(* IEC 61131-3 sources: plc-hackathon-2026/work/dump/MyController/Plc Logic/Application/Init (part 2) *)

(* ---- Init_Prof_FEC.st ---- *)
FUNCTION_BLOCK Init_Prof_FEC
VAR_INPUT
END_VAR
VAR_OUTPUT
END_VAR
VAR
END_VAR

// ---IMPL---
// Inicijalizacija GVL "Prof_FEC"
   Prof_FEC.Data[0] := 40.266;
   Prof_FEC.Data[1] := 42.108;
   Prof_FEC.Data[2] := 42.44;
   Prof_FEC.Data[3] := 43.126;
   Prof_FEC.Data[4] := 43.213;
   Prof_FEC.Data[5] := 42.172;
   Prof_FEC.Data[6] := 44.978;
   Prof_FEC.Data[7] := 44.952;
   Prof_FEC.Data[8] := 43.73;
   Prof_FEC.Data[9] := 41.671;
   Prof_FEC.Data[10] := 39.025;
   Prof_FEC.Data[11] := 43.815;
   Prof_FEC.Data[12] := 42.205;
   Prof_FEC.Data[13] := 42.881;
   Prof_FEC.Data[14] := 40.68;
   Prof_FEC.Data[15] := 39.411;
   Prof_FEC.Data[16] := 40.682;
   Prof_FEC.Data[17] := 40.404;
   Prof_FEC.Data[18] := 41.293;
   Prof_FEC.Data[19] := 41.787;
   Prof_FEC.Data[20] := 254.21;
   Prof_FEC.Data[21] := 268.75;
   Prof_FEC.Data[22] := 265.48;
   Prof_FEC.Data[23] := 296.02;
   Prof_FEC.Data[24] := 335.71;
   Prof_FEC.Data[25] := 339.43;
   Prof_FEC.Data[26] := 388.16;
   Prof_FEC.Data[27] := 433.83;
   Prof_FEC.Data[28] := 441.67;
   Prof_FEC.Data[29] := 486.31;
   Prof_FEC.Data[30] := 552.6;
   Prof_FEC.Data[31] := 544.94;
   Prof_FEC.Data[32] := 568.79;
   Prof_FEC.Data[33] := 634.46;
   Prof_FEC.Data[34] := 604.12;
   Prof_FEC.Data[35] := 630.85;
   Prof_FEC.Data[36] := 656.31;
   Prof_FEC.Data[37] := 671.59;
   Prof_FEC.Data[38] := 634.52;
   Prof_FEC.Data[39] := 653.7;
   Prof_FEC.Data[40] := 625.93;
   Prof_FEC.Data[41] := 654.27;
   Prof_FEC.Data[42] := 603.66;
   Prof_FEC.Data[43] := 590.51;
   Prof_FEC.Data[44] := 620.11;
   Prof_FEC.Data[45] := 604.33;
   Prof_FEC.Data[46] := 589.58;
   Prof_FEC.Data[47] := 638.77;
   Prof_FEC.Data[48] := 571.87;
   Prof_FEC.Data[49] := 540.78;
   Prof_FEC.Data[50] := 589.62;
   Prof_FEC.Data[51] := 576.36;
   Prof_FEC.Data[52] := 646.42;
   Prof_FEC.Data[53] := 628.77;
   Prof_FEC.Data[54] := 633.92;
   Prof_FEC.Data[55] := 671.67;
   Prof_FEC.Data[56] := 731.0;
   Prof_FEC.Data[57] := 742.29;
   Prof_FEC.Data[58] := 722.04;
   Prof_FEC.Data[59] := 711.5;
   Prof_FEC.Data[60] := 722.32;
   Prof_FEC.Data[61] := 679.4;
   Prof_FEC.Data[62] := 676.24;
   Prof_FEC.Data[63] := 745.59;
   Prof_FEC.Data[64] := 789.69;
   Prof_FEC.Data[65] := 795.4;
   Prof_FEC.Data[66] := 766.74;
   Prof_FEC.Data[67] := 673.77;
   Prof_FEC.Data[68] := 501.09;
   Prof_FEC.Data[69] := 365.1;
   Prof_FEC.Data[70] := 325.78;
   Prof_FEC.Data[71] := 293.7;
   Prof_FEC.Data[72] := 276.68;
   Prof_FEC.Data[73] := 266.17;
   Prof_FEC.Data[74] := 227.53;
   Prof_FEC.Data[75] := 256.11;
   Prof_FEC.Data[76] := 43.481;
   Prof_FEC.Data[77] := 44.002;
   Prof_FEC.Data[78] := 44.238;
   Prof_FEC.Data[79] := 43.218;
   Prof_FEC.Data[80] := 40.422;
   Prof_FEC.Data[81] := 41.151;
   Prof_FEC.Data[82] := 40.95;
   Prof_FEC.Data[83] := 41.165;
   Prof_FEC.Data[84] := 40.77;
   Prof_FEC.Data[85] := 43.799;
   Prof_FEC.Data[86] := 42.671;
   Prof_FEC.Data[87] := 43.676;
   Prof_FEC.Data[88] := 41.656;
   Prof_FEC.Data[89] := 40.912;
   Prof_FEC.Data[90] := 41.266;
   Prof_FEC.Data[91] := 39.497;
   Prof_FEC.Data[92] := 44.511;
   Prof_FEC.Data[93] := 44.6;
   Prof_FEC.Data[94] := 47.837;
   Prof_FEC.Data[95] := 45.96;
   Prof_FEC.Data[96] := 45.749;
   Prof_FEC.Data[97] := 44.326;
   Prof_FEC.Data[98] := 44.02;
   Prof_FEC.Data[99] := 43.86;
   Prof_FEC.Data[100] := 44.651;
   Prof_FEC.Data[101] := 48.206;
   Prof_FEC.Data[102] := 43.013;
   Prof_FEC.Data[103] := 45.661;
   Prof_FEC.Data[104] := 40.107;
   Prof_FEC.Data[105] := 41.976;
   Prof_FEC.Data[106] := 37.462;
   Prof_FEC.Data[107] := 40.495;
   Prof_FEC.Data[108] := 45.365;
   Prof_FEC.Data[109] := 47.462;
   Prof_FEC.Data[110] := 48.015;
   Prof_FEC.Data[111] := 48.333;
   Prof_FEC.Data[112] := 47.113;
   Prof_FEC.Data[113] := 48.016;
   Prof_FEC.Data[114] := 44.19;
   Prof_FEC.Data[115] := 45.094;
   Prof_FEC.Data[116] := 290.32;
   Prof_FEC.Data[117] := 297.39;
   Prof_FEC.Data[118] := 284.58;
   Prof_FEC.Data[119] := 325.31;
   Prof_FEC.Data[120] := 357.24;
   Prof_FEC.Data[121] := 394.59;
   Prof_FEC.Data[122] := 407.32;
   Prof_FEC.Data[123] := 458.08;
   Prof_FEC.Data[124] := 551.82;
   Prof_FEC.Data[125] := 580.15;
   Prof_FEC.Data[126] := 608.06;
   Prof_FEC.Data[127] := 578.6;
   Prof_FEC.Data[128] := 612.98;
   Prof_FEC.Data[129] := 614.51;
   Prof_FEC.Data[130] := 640.99;
   Prof_FEC.Data[131] := 677.4;
   Prof_FEC.Data[132] := 743.46;
   Prof_FEC.Data[133] := 772.07;
   Prof_FEC.Data[134] := 790.32;
   Prof_FEC.Data[135] := 764.21;
   Prof_FEC.Data[136] := 693.38;
   Prof_FEC.Data[137] := 715.42;
   Prof_FEC.Data[138] := 590.75;
   Prof_FEC.Data[139] := 678.98;
   Prof_FEC.Data[140] := 643.33;
   Prof_FEC.Data[141] := 614.71;
   Prof_FEC.Data[142] := 677.61;
   Prof_FEC.Data[143] := 646.57;
   Prof_FEC.Data[144] := 662.01;
   Prof_FEC.Data[145] := 656.44;
   Prof_FEC.Data[146] := 583.37;
   Prof_FEC.Data[147] := 664.52;
   Prof_FEC.Data[148] := 554.65;
   Prof_FEC.Data[149] := 629.64;
   Prof_FEC.Data[150] := 670.62;
   Prof_FEC.Data[151] := 596.51;
   Prof_FEC.Data[152] := 661.81;
   Prof_FEC.Data[153] := 592.39;
   Prof_FEC.Data[154] := 608.2;
   Prof_FEC.Data[155] := 668.41;
   Prof_FEC.Data[156] := 618.77;
   Prof_FEC.Data[157] := 575.67;
   Prof_FEC.Data[158] := 513.16;
   Prof_FEC.Data[159] := 598.3;
   Prof_FEC.Data[160] := 660.23;
   Prof_FEC.Data[161] := 656.71;
   Prof_FEC.Data[162] := 634.91;
   Prof_FEC.Data[163] := 512.09;
   Prof_FEC.Data[164] := 414.01;
   Prof_FEC.Data[165] := 373.69;
   Prof_FEC.Data[166] := 339.29;
   Prof_FEC.Data[167] := 286.59;
   Prof_FEC.Data[168] := 285.53;
   Prof_FEC.Data[169] := 218.56;
   Prof_FEC.Data[170] := 242.09;
   Prof_FEC.Data[171] := 257.24;
   Prof_FEC.Data[172] := 44.634;
   Prof_FEC.Data[173] := 44.75;
   Prof_FEC.Data[174] := 41.675;
   Prof_FEC.Data[175] := 49.065;
   Prof_FEC.Data[176] := 47.236;
   Prof_FEC.Data[177] := 43.529;
   Prof_FEC.Data[178] := 44.439;
   Prof_FEC.Data[179] := 44.502;
   Prof_FEC.Data[180] := 48.851;
   Prof_FEC.Data[181] := 50.0;
   Prof_FEC.Data[182] := 47.07;
   Prof_FEC.Data[183] := 44.555;
   Prof_FEC.Data[184] := 44.815;
   Prof_FEC.Data[185] := 44.276;
   Prof_FEC.Data[186] := 44.342;
   Prof_FEC.Data[187] := 43.996;
   Prof_FEC.Data[188] := 44.701;
   Prof_FEC.Data[189] := 45.391;
   Prof_FEC.Data[190] := 41.212;
   Prof_FEC.Data[191] := 44.161;
   Prof_FEC.Data[192] := 43.203;
   Prof_FEC.Data[193] := 41.683;
   Prof_FEC.Data[194] := 43.808;
   Prof_FEC.Data[195] := 42.414;
   Prof_FEC.Data[196] := 40.31;
   Prof_FEC.Data[197] := 46.212;
   Prof_FEC.Data[198] := 49.298;
   Prof_FEC.Data[199] := 47.323;
   Prof_FEC.Data[200] := 45.775;
   Prof_FEC.Data[201] := 44.057;
   Prof_FEC.Data[202] := 46.892;
   Prof_FEC.Data[203] := 46.929;
   Prof_FEC.Data[204] := 47.35;
   Prof_FEC.Data[205] := 50.0;
   Prof_FEC.Data[206] := 49.345;
   Prof_FEC.Data[207] := 45.771;
   Prof_FEC.Data[208] := 45.917;
   Prof_FEC.Data[209] := 42.603;
   Prof_FEC.Data[210] := 42.491;
   Prof_FEC.Data[211] := 45.313;
   Prof_FEC.Data[212] := 319.06;
   Prof_FEC.Data[213] := 330.88;
   Prof_FEC.Data[214] := 322.58;
   Prof_FEC.Data[215] := 340.34;
   Prof_FEC.Data[216] := 275.1;
   Prof_FEC.Data[217] := 281.37;
   Prof_FEC.Data[218] := 266.89;
   Prof_FEC.Data[219] := 303.74;
   Prof_FEC.Data[220] := 373.21;
   Prof_FEC.Data[221] := 357.72;
   Prof_FEC.Data[222] := 340.19;
   Prof_FEC.Data[223] := 329.95;
   Prof_FEC.Data[224] := 295.08;
   Prof_FEC.Data[225] := 279.44;
   Prof_FEC.Data[226] := 275.77;
   Prof_FEC.Data[227] := 307.14;
   Prof_FEC.Data[228] := 325.7;
   Prof_FEC.Data[229] := 380.71;
   Prof_FEC.Data[230] := 366.07;
   Prof_FEC.Data[231] := 385.12;
   Prof_FEC.Data[232] := 384.91;
   Prof_FEC.Data[233] := 335.32;
   Prof_FEC.Data[234] := 372.66;
   Prof_FEC.Data[235] := 336.27;
   Prof_FEC.Data[236] := 358.41;
   Prof_FEC.Data[237] := 372.35;
   Prof_FEC.Data[238] := 376.62;
   Prof_FEC.Data[239] := 316.95;
   Prof_FEC.Data[240] := 316.07;
   Prof_FEC.Data[241] := 285.92;
   Prof_FEC.Data[242] := 287.26;
   Prof_FEC.Data[243] := 332.84;
   Prof_FEC.Data[244] := 301.17;
   Prof_FEC.Data[245] := 295.5;
   Prof_FEC.Data[246] := 302.52;
   Prof_FEC.Data[247] := 302.02;
   Prof_FEC.Data[248] := 289.77;
   Prof_FEC.Data[249] := 294.29;
   Prof_FEC.Data[250] := 289.81;
   Prof_FEC.Data[251] := 281.9;
   Prof_FEC.Data[252] := 305.51;
   Prof_FEC.Data[253] := 338.99;
   Prof_FEC.Data[254] := 298.04;
   Prof_FEC.Data[255] := 304.85;
   Prof_FEC.Data[256] := 262.63;
   Prof_FEC.Data[257] := 289.06;
   Prof_FEC.Data[258] := 310.2;
   Prof_FEC.Data[259] := 302.52;
   Prof_FEC.Data[260] := 297.0;
   Prof_FEC.Data[261] := 316.44;
   Prof_FEC.Data[262] := 313.22;
   Prof_FEC.Data[263] := 331.56;
   Prof_FEC.Data[264] := 356.25;
   Prof_FEC.Data[265] := 332.19;
   Prof_FEC.Data[266] := 338.85;
   Prof_FEC.Data[267] := 311.86;
   Prof_FEC.Data[268] := 43.718;
   Prof_FEC.Data[269] := 41.336;
   Prof_FEC.Data[270] := 42.442;
   Prof_FEC.Data[271] := 43.645;
   Prof_FEC.Data[272] := 46.923;
   Prof_FEC.Data[273] := 47.891;
   Prof_FEC.Data[274] := 47.964;
   Prof_FEC.Data[275] := 49.914;
   Prof_FEC.Data[276] := 44.567;
   Prof_FEC.Data[277] := 40.108;
   Prof_FEC.Data[278] := 42.664;
   Prof_FEC.Data[279] := 42.486;
   Prof_FEC.Data[280] := 44.943;
   Prof_FEC.Data[281] := 50.0;
   Prof_FEC.Data[282] := 50.0;
   Prof_FEC.Data[283] := 47.638;
   Prof_FEC.Data[284] := 50.0;
   Prof_FEC.Data[285] := 49.774;
   Prof_FEC.Data[286] := 48.766;
   Prof_FEC.Data[287] := 49.774;
   Prof_FEC.Data[288] := 49.582;
   Prof_FEC.Data[289] := 50.0;
   Prof_FEC.Data[290] := 50.0;
   Prof_FEC.Data[291] := 50.0;
   Prof_FEC.Data[292] := 47.656;
   Prof_FEC.Data[293] := 45.649;
   Prof_FEC.Data[294] := 47.716;
   Prof_FEC.Data[295] := 47.822;
   Prof_FEC.Data[296] := 50.0;
   Prof_FEC.Data[297] := 50.0;
   Prof_FEC.Data[298] := 50.0;
   Prof_FEC.Data[299] := 50.0;
   Prof_FEC.Data[300] := 49.981;
   Prof_FEC.Data[301] := 42.622;
   Prof_FEC.Data[302] := 45.328;
   Prof_FEC.Data[303] := 41.662;
   Prof_FEC.Data[304] := 42.786;
   Prof_FEC.Data[305] := 46.932;
   Prof_FEC.Data[306] := 47.834;
   Prof_FEC.Data[307] := 46.461;
   Prof_FEC.Data[308] := 283.9;
   Prof_FEC.Data[309] := 312.44;
   Prof_FEC.Data[310] := 294.91;
   Prof_FEC.Data[311] := 326.05;
   Prof_FEC.Data[312] := 357.35;
   Prof_FEC.Data[313] := 376.04;
   Prof_FEC.Data[314] := 408.97;
   Prof_FEC.Data[315] := 349.34;
   Prof_FEC.Data[316] := 322.6;
   Prof_FEC.Data[317] := 310.61;
   Prof_FEC.Data[318] := 331.18;
   Prof_FEC.Data[319] := 318.25;
   Prof_FEC.Data[320] := 269.4;
   Prof_FEC.Data[321] := 240.37;
   Prof_FEC.Data[322] := 213.63;
   Prof_FEC.Data[323] := 225.18;
   Prof_FEC.Data[324] := 185.0;
   Prof_FEC.Data[325] := 166.18;
   Prof_FEC.Data[326] := 187.61;
   Prof_FEC.Data[327] := 197.79;
   Prof_FEC.Data[328] := 225.46;
   Prof_FEC.Data[329] := 225.06;
   Prof_FEC.Data[330] := 228.64;
   Prof_FEC.Data[331] := 195.52;
   Prof_FEC.Data[332] := 174.06;
   Prof_FEC.Data[333] := 170.88;
   Prof_FEC.Data[334] := 175.29;
   Prof_FEC.Data[335] := 215.34;
   Prof_FEC.Data[336] := 203.35;
   Prof_FEC.Data[337] := 211.31;
   Prof_FEC.Data[338] := 223.33;
   Prof_FEC.Data[339] := 212.28;
   Prof_FEC.Data[340] := 167.16;
   Prof_FEC.Data[341] := 183.77;
   Prof_FEC.Data[342] := 163.03;
   Prof_FEC.Data[343] := 134.03;
   Prof_FEC.Data[344] := 177.4;
   Prof_FEC.Data[345] := 184.68;
   Prof_FEC.Data[346] := 189.82;
   Prof_FEC.Data[347] := 188.48;
   Prof_FEC.Data[348] := 164.02;
   Prof_FEC.Data[349] := 156.08;
   Prof_FEC.Data[350] := 174.91;
   Prof_FEC.Data[351] := 205.13;
   Prof_FEC.Data[352] := 252.54;
   Prof_FEC.Data[353] := 249.88;
   Prof_FEC.Data[354] := 261.78;
   Prof_FEC.Data[355] := 335.45;
   Prof_FEC.Data[356] := 293.76;
   Prof_FEC.Data[357] := 307.86;
   Prof_FEC.Data[358] := 290.99;
   Prof_FEC.Data[359] := 264.47;
   Prof_FEC.Data[360] := 300.89;
   Prof_FEC.Data[361] := 319.15;
   Prof_FEC.Data[362] := 295.24;
   Prof_FEC.Data[363] := 350.74;
   Prof_FEC.Data[364] := 44.223;
   Prof_FEC.Data[365] := 43.602;
   Prof_FEC.Data[366] := 42.21;
   Prof_FEC.Data[367] := 49.285;
   Prof_FEC.Data[368] := 50.0;
   Prof_FEC.Data[369] := 50.0;
   Prof_FEC.Data[370] := 50.0;
   Prof_FEC.Data[371] := 49.043;
   Prof_FEC.Data[372] := 47.995;
   Prof_FEC.Data[373] := 46.41;
   Prof_FEC.Data[374] := 45.867;
   Prof_FEC.Data[375] := 47.788;
   Prof_FEC.Data[376] := 50.0;
   Prof_FEC.Data[377] := 50.0;
   Prof_FEC.Data[378] := 50.0;
   Prof_FEC.Data[379] := 49.985;
   Prof_FEC.Data[380] := 47.547;
   Prof_FEC.Data[381] := 47.572;
   Prof_FEC.Data[382] := 48.112;
   Prof_FEC.Data[383] := 48.506;
   Prof_FEC.Data[384] := 41.761;
   Prof_FEC.Data[385] := 40.506;
   Prof_FEC.Data[386] := 41.058;
   Prof_FEC.Data[387] := 41.3;
   Prof_FEC.Data[388] := 37.893;
   Prof_FEC.Data[389] := 36.404;
   Prof_FEC.Data[390] := 39.255;
   Prof_FEC.Data[391] := 39.306;
   Prof_FEC.Data[392] := 39.088;
   Prof_FEC.Data[393] := 41.274;
   Prof_FEC.Data[394] := 41.431;
   Prof_FEC.Data[395] := 40.833;
   Prof_FEC.Data[396] := 38.292;
   Prof_FEC.Data[397] := 40.541;
   Prof_FEC.Data[398] := 42.673;
   Prof_FEC.Data[399] := 40.341;
   Prof_FEC.Data[400] := 43.559;
   Prof_FEC.Data[401] := 41.749;
   Prof_FEC.Data[402] := 44.034;
   Prof_FEC.Data[403] := 42.021;
   Prof_FEC.Data[404] := 220.86;
   Prof_FEC.Data[405] := 231.61;
   Prof_FEC.Data[406] := 252.32;
   Prof_FEC.Data[407] := 268.96;
   Prof_FEC.Data[408] := 267.93;
   Prof_FEC.Data[409] := 273.79;
   Prof_FEC.Data[410] := 270.15;
   Prof_FEC.Data[411] := 295.92;
   Prof_FEC.Data[412] := 295.59;
   Prof_FEC.Data[413] := 262.91;
   Prof_FEC.Data[414] := 252.04;
   Prof_FEC.Data[415] := 217.69;
   Prof_FEC.Data[416] := 191.04;
   Prof_FEC.Data[417] := 157.39;
   Prof_FEC.Data[418] := 138.36;
   Prof_FEC.Data[419] := 143.73;
   Prof_FEC.Data[420] := 129.02;
   Prof_FEC.Data[421] := 131.7;
   Prof_FEC.Data[422] := 120.58;
   Prof_FEC.Data[423] := 123.58;
   Prof_FEC.Data[424] := 147.65;
   Prof_FEC.Data[425] := 154.92;
   Prof_FEC.Data[426] := 156.45;
   Prof_FEC.Data[427] := 156.39;
   Prof_FEC.Data[428] := 137.58;
   Prof_FEC.Data[429] := 126.17;
   Prof_FEC.Data[430] := 126.61;
   Prof_FEC.Data[431] := 129.68;
   Prof_FEC.Data[432] := 140.12;
   Prof_FEC.Data[433] := 157.56;
   Prof_FEC.Data[434] := 151.75;
   Prof_FEC.Data[435] := 162.25;
   Prof_FEC.Data[436] := 128.1;
   Prof_FEC.Data[437] := 126.78;
   Prof_FEC.Data[438] := 117.5;
   Prof_FEC.Data[439] := 118.93;
   Prof_FEC.Data[440] := 142.47;
   Prof_FEC.Data[441] := 152.95;
   Prof_FEC.Data[442] := 149.14;
   Prof_FEC.Data[443] := 145.03;
   Prof_FEC.Data[444] := 117.79;
   Prof_FEC.Data[445] := 111.38;
   Prof_FEC.Data[446] := 104.69;
   Prof_FEC.Data[447] := 141.73;
   Prof_FEC.Data[448] := 212.13;
   Prof_FEC.Data[449] := 224.04;
   Prof_FEC.Data[450] := 228.65;
   Prof_FEC.Data[451] := 248.51;
   Prof_FEC.Data[452] := 255.06;
   Prof_FEC.Data[453] := 245.97;
   Prof_FEC.Data[454] := 262.91;
   Prof_FEC.Data[455] := 267.76;
   Prof_FEC.Data[456] := 223.68;
   Prof_FEC.Data[457] := 256.21;
   Prof_FEC.Data[458] := 232.8;
   Prof_FEC.Data[459] := 274.8;
   Prof_FEC.Data[460] := 39.079;
   Prof_FEC.Data[461] := 39.025;
   Prof_FEC.Data[462] := 41.564;
   Prof_FEC.Data[463] := 38.951;
   Prof_FEC.Data[464] := 40.754;
   Prof_FEC.Data[465] := 39.858;
   Prof_FEC.Data[466] := 44.481;
   Prof_FEC.Data[467] := 43.308;
   Prof_FEC.Data[468] := 38.958;
   Prof_FEC.Data[469] := 37.768;
   Prof_FEC.Data[470] := 40.13;
   Prof_FEC.Data[471] := 43.311;
   Prof_FEC.Data[472] := 41.868;
   Prof_FEC.Data[473] := 41.644;
   Prof_FEC.Data[474] := 45.684;
   Prof_FEC.Data[475] := 41.713;
   Prof_FEC.Data[476] := 40.566;
   Prof_FEC.Data[477] := 37.16;
   Prof_FEC.Data[478] := 38.8;
   Prof_FEC.Data[479] := 37.164;
   Prof_FEC.Data[480] := 41.382;
   Prof_FEC.Data[481] := 38.333;
   Prof_FEC.Data[482] := 41.534;
   Prof_FEC.Data[483] := 39.258;
   Prof_FEC.Data[484] := 37.921;
   Prof_FEC.Data[485] := 39.211;
   Prof_FEC.Data[486] := 38.448;
   Prof_FEC.Data[487] := 39.102;
   Prof_FEC.Data[488] := 40.047;
   Prof_FEC.Data[489] := 42.576;
   Prof_FEC.Data[490] := 38.555;
   Prof_FEC.Data[491] := 42.984;
   Prof_FEC.Data[492] := 39.987;
   Prof_FEC.Data[493] := 37.635;
   Prof_FEC.Data[494] := 39.065;
   Prof_FEC.Data[495] := 39.048;
   Prof_FEC.Data[496] := 41.244;
   Prof_FEC.Data[497] := 39.491;
   Prof_FEC.Data[498] := 42.125;
   Prof_FEC.Data[499] := 40.701;
   Prof_FEC.Data[500] := 233.19;
   Prof_FEC.Data[501] := 246.58;
   Prof_FEC.Data[502] := 243.83;
   Prof_FEC.Data[503] := 281.26;
   Prof_FEC.Data[504] := 295.39;
   Prof_FEC.Data[505] := 370.32;
   Prof_FEC.Data[506] := 397.69;
   Prof_FEC.Data[507] := 455.67;
   Prof_FEC.Data[508] := 520.44;
   Prof_FEC.Data[509] := 553.71;
   Prof_FEC.Data[510] := 689.15;
   Prof_FEC.Data[511] := 598.67;
   Prof_FEC.Data[512] := 572.27;
   Prof_FEC.Data[513] := 519.77;
   Prof_FEC.Data[514] := 583.63;
   Prof_FEC.Data[515] := 549.88;
   Prof_FEC.Data[516] := 620.15;
   Prof_FEC.Data[517] := 653.48;
   Prof_FEC.Data[518] := 602.24;
   Prof_FEC.Data[519] := 566.8;
   Prof_FEC.Data[520] := 516.28;
   Prof_FEC.Data[521] := 602.42;
   Prof_FEC.Data[522] := 637.19;
   Prof_FEC.Data[523] := 681.85;
   Prof_FEC.Data[524] := 777.61;
   Prof_FEC.Data[525] := 736.14;
   Prof_FEC.Data[526] := 590.05;
   Prof_FEC.Data[527] := 649.37;
   Prof_FEC.Data[528] := 574.35;
   Prof_FEC.Data[529] := 592.82;
   Prof_FEC.Data[530] := 547.79;
   Prof_FEC.Data[531] := 566.16;
   Prof_FEC.Data[532] := 665.87;
   Prof_FEC.Data[533] := 677.43;
   Prof_FEC.Data[534] := 703.62;
   Prof_FEC.Data[535] := 625.62;
   Prof_FEC.Data[536] := 547.25;
   Prof_FEC.Data[537] := 620.27;
   Prof_FEC.Data[538] := 624.7;
   Prof_FEC.Data[539] := 656.31;
   Prof_FEC.Data[540] := 606.26;
   Prof_FEC.Data[541] := 616.95;
   Prof_FEC.Data[542] := 668.6;
   Prof_FEC.Data[543] := 616.15;
   Prof_FEC.Data[544] := 698.59;
   Prof_FEC.Data[545] := 831.84;
   Prof_FEC.Data[546] := 817.44;
   Prof_FEC.Data[547] := 650.21;
   Prof_FEC.Data[548] := 449.5;
   Prof_FEC.Data[549] := 357.2;
   Prof_FEC.Data[550] := 340.66;
   Prof_FEC.Data[551] := 329.73;
   Prof_FEC.Data[552] := 276.28;
   Prof_FEC.Data[553] := 251.0;
   Prof_FEC.Data[554] := 243.4;
   Prof_FEC.Data[555] := 235.76;
   Prof_FEC.Data[556] := 41.455;
   Prof_FEC.Data[557] := 41.369;
   Prof_FEC.Data[558] := 42.919;
   Prof_FEC.Data[559] := 42.389;
   Prof_FEC.Data[560] := 43.311;
   Prof_FEC.Data[561] := 39.254;
   Prof_FEC.Data[562] := 39.57;
   Prof_FEC.Data[563] := 43.124;
   Prof_FEC.Data[564] := 44.513;
   Prof_FEC.Data[565] := 45.492;
   Prof_FEC.Data[566] := 47.736;
   Prof_FEC.Data[567] := 45.711;
   Prof_FEC.Data[568] := 44.029;
   Prof_FEC.Data[569] := 44.732;
   Prof_FEC.Data[570] := 44.758;
   Prof_FEC.Data[571] := 45.416;
   Prof_FEC.Data[572] := 43.543;
   Prof_FEC.Data[573] := 47.234;
   Prof_FEC.Data[574] := 50.0;
   Prof_FEC.Data[575] := 50.0;
   Prof_FEC.Data[576] := 43.237;
   Prof_FEC.Data[577] := 45.836;
   Prof_FEC.Data[578] := 44.0;
   Prof_FEC.Data[579] := 43.91;
   Prof_FEC.Data[580] := 45.488;
   Prof_FEC.Data[581] := 47.976;
   Prof_FEC.Data[582] := 47.802;
   Prof_FEC.Data[583] := 49.458;
   Prof_FEC.Data[584] := 42.187;
   Prof_FEC.Data[585] := 42.069;
   Prof_FEC.Data[586] := 46.957;
   Prof_FEC.Data[587] := 45.27;
   Prof_FEC.Data[588] := 44.793;
   Prof_FEC.Data[589] := 46.33;
   Prof_FEC.Data[590] := 43.176;
   Prof_FEC.Data[591] := 44.03;
   Prof_FEC.Data[592] := 40.855;
   Prof_FEC.Data[593] := 41.644;
   Prof_FEC.Data[594] := 42.269;
   Prof_FEC.Data[595] := 41.999;
   Prof_FEC.Data[596] := 263.51;
   Prof_FEC.Data[597] := 287.36;
   Prof_FEC.Data[598] := 286.34;
   Prof_FEC.Data[599] := 304.23;
   Prof_FEC.Data[600] := 335.11;
   Prof_FEC.Data[601] := 377.91;
   Prof_FEC.Data[602] := 432.91;
   Prof_FEC.Data[603] := 417.93;
   Prof_FEC.Data[604] := 508.5;
   Prof_FEC.Data[605] := 524.9;
   Prof_FEC.Data[606] := 537.3;
   Prof_FEC.Data[607] := 526.95;
   Prof_FEC.Data[608] := 541.55;
   Prof_FEC.Data[609] := 573.71;
   Prof_FEC.Data[610] := 591.4;
   Prof_FEC.Data[611] := 602.76;
   Prof_FEC.Data[612] := 785.56;
   Prof_FEC.Data[613] := 734.56;
   Prof_FEC.Data[614] := 706.14;
   Prof_FEC.Data[615] := 716.39;
   Prof_FEC.Data[616] := 661.63;
   Prof_FEC.Data[617] := 678.87;
   Prof_FEC.Data[618] := 710.72;
   Prof_FEC.Data[619] := 696.29;
   Prof_FEC.Data[620] := 634.02;
   Prof_FEC.Data[621] := 643.44;
   Prof_FEC.Data[622] := 550.0;
   Prof_FEC.Data[623] := 566.25;
   Prof_FEC.Data[624] := 589.4;
   Prof_FEC.Data[625] := 555.62;
   Prof_FEC.Data[626] := 459.68;
   Prof_FEC.Data[627] := 476.96;
   Prof_FEC.Data[628] := 619.81;
   Prof_FEC.Data[629] := 575.1;
   Prof_FEC.Data[630] := 556.24;
   Prof_FEC.Data[631] := 604.41;
   Prof_FEC.Data[632] := 654.33;
   Prof_FEC.Data[633] := 615.72;
   Prof_FEC.Data[634] := 599.9;
   Prof_FEC.Data[635] := 669.87;
   Prof_FEC.Data[636] := 671.34;
   Prof_FEC.Data[637] := 665.18;
   Prof_FEC.Data[638] := 665.52;
   Prof_FEC.Data[639] := 732.21;
   Prof_FEC.Data[640] := 802.07;
   Prof_FEC.Data[641] := 828.81;
   Prof_FEC.Data[642] := 759.3;
   Prof_FEC.Data[643] := 593.23;
   Prof_FEC.Data[644] := 440.78;
   Prof_FEC.Data[645] := 373.82;
   Prof_FEC.Data[646] := 324.14;
   Prof_FEC.Data[647] := 305.19;
   Prof_FEC.Data[648] := 261.91;
   Prof_FEC.Data[649] := 253.88;
   Prof_FEC.Data[650] := 240.22;
   Prof_FEC.Data[651] := 270.32;
   Prof_FEC.Data[652] := 43.725;
   Prof_FEC.Data[653] := 44.364;
   Prof_FEC.Data[654] := 43.17;
   Prof_FEC.Data[655] := 42.668;
   Prof_FEC.Data[656] := 39.396;
   Prof_FEC.Data[657] := 40.766;
   Prof_FEC.Data[658] := 43.679;
   Prof_FEC.Data[659] := 44.295;
   Prof_FEC.Data[660] := 45.57;
   Prof_FEC.Data[661] := 46.176;
   Prof_FEC.Data[662] := 46.012;
   Prof_FEC.Data[663] := 44.906;
   Prof_FEC.Data[664] := 43.523;
   Prof_FEC.Data[665] := 42.009;
   Prof_FEC.Data[666] := 41.989;
   Prof_FEC.Data[667] := 44.79;
   Prof_FEC.Data[668] := 44.326;
   Prof_FEC.Data[669] := 44.936;
   Prof_FEC.Data[670] := 43.69;
   Prof_FEC.Data[671] := 45.738;
   Prof_FEC.Data[672] := 44.028;
   Prof_FEC.Data[673] := 39.767;
   Prof_FEC.Data[674] := 41.813;
   Prof_FEC.Data[675] := 41.887;
   Prof_FEC.Data[676] := 45.51;
   Prof_FEC.Data[677] := 44.014;
   Prof_FEC.Data[678] := 40.069;
   Prof_FEC.Data[679] := 43.938;
   Prof_FEC.Data[680] := 42.852;
   Prof_FEC.Data[681] := 42.118;
   Prof_FEC.Data[682] := 38.044;
   Prof_FEC.Data[683] := 40.184;
   Prof_FEC.Data[684] := 42.822;
   Prof_FEC.Data[685] := 40.133;
   Prof_FEC.Data[686] := 42.875;
   Prof_FEC.Data[687] := 41.446;
   Prof_FEC.Data[688] := 41.683;
   Prof_FEC.Data[689] := 37.861;
   Prof_FEC.Data[690] := 38.58;
   Prof_FEC.Data[691] := 40.941;
   Prof_FEC.Data[692] := 282.48;
   Prof_FEC.Data[693] := 332.35;
   Prof_FEC.Data[694] := 325.29;
   Prof_FEC.Data[695] := 335.58;
   Prof_FEC.Data[696] := 395.27;
   Prof_FEC.Data[697] := 452.43;
   Prof_FEC.Data[698] := 454.87;
   Prof_FEC.Data[699] := 541.36;
   Prof_FEC.Data[700] := 585.95;
   Prof_FEC.Data[701] := 601.86;
   Prof_FEC.Data[702] := 594.43;
   Prof_FEC.Data[703] := 648.13;
   Prof_FEC.Data[704] := 588.8;
   Prof_FEC.Data[705] := 612.08;
   Prof_FEC.Data[706] := 634.29;
   Prof_FEC.Data[707] := 622.98;
   Prof_FEC.Data[708] := 736.64;
   Prof_FEC.Data[709] := 734.86;
   Prof_FEC.Data[710] := 722.76;
   Prof_FEC.Data[711] := 751.4;
   Prof_FEC.Data[712] := 718.86;
   Prof_FEC.Data[713] := 681.41;
   Prof_FEC.Data[714] := 682.09;
   Prof_FEC.Data[715] := 698.66;
   Prof_FEC.Data[716] := 684.77;
   Prof_FEC.Data[717] := 611.4;
   Prof_FEC.Data[718] := 677.7;
   Prof_FEC.Data[719] := 583.36;
   Prof_FEC.Data[720] := 598.17;
   Prof_FEC.Data[721] := 548.09;
   Prof_FEC.Data[722] := 578.6;
   Prof_FEC.Data[723] := 658.22;
   Prof_FEC.Data[724] := 620.59;
   Prof_FEC.Data[725] := 577.57;
   Prof_FEC.Data[726] := 629.63;
   Prof_FEC.Data[727] := 666.61;
   Prof_FEC.Data[728] := 665.39;
   Prof_FEC.Data[729] := 629.68;
   Prof_FEC.Data[730] := 638.08;
   Prof_FEC.Data[731] := 645.85;
   Prof_FEC.Data[732] := 571.4;
   Prof_FEC.Data[733] := 637.63;
   Prof_FEC.Data[734] := 645.71;
   Prof_FEC.Data[735] := 751.55;
   Prof_FEC.Data[736] := 766.08;
   Prof_FEC.Data[737] := 817.3;
   Prof_FEC.Data[738] := 804.18;
   Prof_FEC.Data[739] := 678.1;
   Prof_FEC.Data[740] := 476.49;
   Prof_FEC.Data[741] := 411.55;
   Prof_FEC.Data[742] := 340.04;
   Prof_FEC.Data[743] := 333.82;
   Prof_FEC.Data[744] := 289.65;
   Prof_FEC.Data[745] := 264.09;
   Prof_FEC.Data[746] := 258.98;
   Prof_FEC.Data[747] := 238.7;
   Prof_FEC.Data[748] := 41.003;
   Prof_FEC.Data[749] := 43.086;
   Prof_FEC.Data[750] := 44.613;
   Prof_FEC.Data[751] := 44.27;
   Prof_FEC.Data[752] := 41.883;
   Prof_FEC.Data[753] := 40.89;
   Prof_FEC.Data[754] := 43.059;
   Prof_FEC.Data[755] := 41.991;
   Prof_FEC.Data[756] := 43.288;
   Prof_FEC.Data[757] := 46.229;
   Prof_FEC.Data[758] := 47.842;
   Prof_FEC.Data[759] := 46.058;
   Prof_FEC.Data[760] := 42.668;
   Prof_FEC.Data[761] := 42.378;
   Prof_FEC.Data[762] := 44.29;
   Prof_FEC.Data[763] := 39.668;
   Prof_FEC.Data[764] := 46.148;
   Prof_FEC.Data[765] := 44.498;
   Prof_FEC.Data[766] := 45.658;
   Prof_FEC.Data[767] := 40.353;
   Prof_FEC.Data[768] := 38.277;
   Prof_FEC.Data[769] := 39.793;
   Prof_FEC.Data[770] := 40.946;
   Prof_FEC.Data[771] := 40.44;
   Prof_FEC.Data[772] := 45.389;
   Prof_FEC.Data[773] := 40.252;
   Prof_FEC.Data[774] := 38.412;
   Prof_FEC.Data[775] := 39.232;
   Prof_FEC.Data[776] := 37.656;
   Prof_FEC.Data[777] := 38.556;
   Prof_FEC.Data[778] := 38.034;
   Prof_FEC.Data[779] := 40.356;
   Prof_FEC.Data[780] := 42.612;
   Prof_FEC.Data[781] := 44.846;
   Prof_FEC.Data[782] := 42.507;
   Prof_FEC.Data[783] := 42.493;
   Prof_FEC.Data[784] := 41.157;
   Prof_FEC.Data[785] := 40.099;
   Prof_FEC.Data[786] := 40.519;
   Prof_FEC.Data[787] := 38.419;
   Prof_FEC.Data[788] := 261.11;
   Prof_FEC.Data[789] := 270.77;
   Prof_FEC.Data[790] := 279.01;
   Prof_FEC.Data[791] := 306.17;
   Prof_FEC.Data[792] := 312.74;
   Prof_FEC.Data[793] := 367.39;
   Prof_FEC.Data[794] := 372.22;
   Prof_FEC.Data[795] := 403.09;
   Prof_FEC.Data[796] := 368.48;
   Prof_FEC.Data[797] := 439.71;
   Prof_FEC.Data[798] := 435.87;
   Prof_FEC.Data[799] := 519.7;
   Prof_FEC.Data[800] := 543.18;
   Prof_FEC.Data[801] := 599.16;
   Prof_FEC.Data[802] := 574.9;
   Prof_FEC.Data[803] := 630.27;
   Prof_FEC.Data[804] := 658.4;
   Prof_FEC.Data[805] := 666.64;
   Prof_FEC.Data[806] := 648.09;
   Prof_FEC.Data[807] := 637.81;
   Prof_FEC.Data[808] := 663.44;
   Prof_FEC.Data[809] := 598.05;
   Prof_FEC.Data[810] := 613.49;
   Prof_FEC.Data[811] := 658.19;
   Prof_FEC.Data[812] := 624.31;
   Prof_FEC.Data[813] := 648.27;
   Prof_FEC.Data[814] := 608.76;
   Prof_FEC.Data[815] := 653.53;
   Prof_FEC.Data[816] := 620.42;
   Prof_FEC.Data[817] := 610.22;
   Prof_FEC.Data[818] := 566.41;
   Prof_FEC.Data[819] := 578.15;
   Prof_FEC.Data[820] := 597.42;
   Prof_FEC.Data[821] := 589.31;
   Prof_FEC.Data[822] := 617.84;
   Prof_FEC.Data[823] := 542.02;
   Prof_FEC.Data[824] := 607.11;
   Prof_FEC.Data[825] := 669.5;
   Prof_FEC.Data[826] := 660.41;
   Prof_FEC.Data[827] := 687.15;
   Prof_FEC.Data[828] := 657.45;
   Prof_FEC.Data[829] := 582.33;
   Prof_FEC.Data[830] := 611.92;
   Prof_FEC.Data[831] := 625.45;
   Prof_FEC.Data[832] := 723.16;
   Prof_FEC.Data[833] := 835.76;
   Prof_FEC.Data[834] := 808.77;
   Prof_FEC.Data[835] := 671.07;
   Prof_FEC.Data[836] := 512.07;
   Prof_FEC.Data[837] := 427.59;
   Prof_FEC.Data[838] := 364.39;
   Prof_FEC.Data[839] := 294.08;
   Prof_FEC.Data[840] := 312.99;
   Prof_FEC.Data[841] := 263.95;
   Prof_FEC.Data[842] := 257.21;
   Prof_FEC.Data[843] := 263.71;
   Prof_FEC.Data[844] := 43.381;
   Prof_FEC.Data[845] := 42.586;
   Prof_FEC.Data[846] := 41.597;
   Prof_FEC.Data[847] := 38.529;
   Prof_FEC.Data[848] := 36.848;
   Prof_FEC.Data[849] := 36.427;
   Prof_FEC.Data[850] := 35.903;
   Prof_FEC.Data[851] := 40.35;
   Prof_FEC.Data[852] := 40.966;
   Prof_FEC.Data[853] := 39.394;
   Prof_FEC.Data[854] := 41.652;
   Prof_FEC.Data[855] := 39.939;
   Prof_FEC.Data[856] := 41.507;
   Prof_FEC.Data[857] := 39.621;
   Prof_FEC.Data[858] := 38.222;
   Prof_FEC.Data[859] := 40.901;
   Prof_FEC.Data[860] := 42.692;
   Prof_FEC.Data[861] := 41.806;
   Prof_FEC.Data[862] := 44.237;
   Prof_FEC.Data[863] := 42.542;
   Prof_FEC.Data[864] := 43.501;
   Prof_FEC.Data[865] := 42.176;
   Prof_FEC.Data[866] := 42.518;
   Prof_FEC.Data[867] := 42.429;
   Prof_FEC.Data[868] := 43.879;
   Prof_FEC.Data[869] := 44.418;
   Prof_FEC.Data[870] := 41.657;
   Prof_FEC.Data[871] := 44.324;
   Prof_FEC.Data[872] := 41.629;
   Prof_FEC.Data[873] := 39.627;
   Prof_FEC.Data[874] := 42.944;
   Prof_FEC.Data[875] := 44.603;
   Prof_FEC.Data[876] := 43.197;
   Prof_FEC.Data[877] := 43.806;
   Prof_FEC.Data[878] := 45.903;
   Prof_FEC.Data[879] := 45.022;
   Prof_FEC.Data[880] := 41.083;
   Prof_FEC.Data[881] := 41.415;
   Prof_FEC.Data[882] := 39.237;
   Prof_FEC.Data[883] := 40.072;
   Prof_FEC.Data[884] := 239.42;
   Prof_FEC.Data[885] := 257.82;
   Prof_FEC.Data[886] := 279.46;
   Prof_FEC.Data[887] := 243.95;
   Prof_FEC.Data[888] := 315.84;
   Prof_FEC.Data[889] := 312.15;
   Prof_FEC.Data[890] := 397.45;
   Prof_FEC.Data[891] := 464.0;
   Prof_FEC.Data[892] := 453.22;
   Prof_FEC.Data[893] := 490.71;
   Prof_FEC.Data[894] := 497.23;
   Prof_FEC.Data[895] := 466.06;
   Prof_FEC.Data[896] := 567.12;
   Prof_FEC.Data[897] := 516.2;
   Prof_FEC.Data[898] := 597.08;
   Prof_FEC.Data[899] := 567.75;
   Prof_FEC.Data[900] := 628.95;
   Prof_FEC.Data[901] := 666.07;
   Prof_FEC.Data[902] := 628.96;
   Prof_FEC.Data[903] := 696.53;
   Prof_FEC.Data[904] := 696.22;
   Prof_FEC.Data[905] := 640.4;
   Prof_FEC.Data[906] := 659.8;
   Prof_FEC.Data[907] := 706.87;
   Prof_FEC.Data[908] := 750.8;
   Prof_FEC.Data[909] := 743.56;
   Prof_FEC.Data[910] := 691.18;
   Prof_FEC.Data[911] := 680.06;
   Prof_FEC.Data[912] := 653.39;
   Prof_FEC.Data[913] := 702.72;
   Prof_FEC.Data[914] := 631.86;
   Prof_FEC.Data[915] := 622.26;
   Prof_FEC.Data[916] := 653.05;
   Prof_FEC.Data[917] := 664.46;
   Prof_FEC.Data[918] := 695.22;
   Prof_FEC.Data[919] := 705.99;
   Prof_FEC.Data[920] := 644.67;
   Prof_FEC.Data[921] := 677.48;
   Prof_FEC.Data[922] := 548.97;
   Prof_FEC.Data[923] := 603.14;
   Prof_FEC.Data[924] := 617.86;
   Prof_FEC.Data[925] := 549.85;
   Prof_FEC.Data[926] := 550.91;
   Prof_FEC.Data[927] := 653.21;
   Prof_FEC.Data[928] := 646.05;
   Prof_FEC.Data[929] := 772.32;
   Prof_FEC.Data[930] := 793.02;
   Prof_FEC.Data[931] := 569.74;
   Prof_FEC.Data[932] := 445.62;
   Prof_FEC.Data[933] := 315.95;
   Prof_FEC.Data[934] := 271.18;
   Prof_FEC.Data[935] := 267.25;
   Prof_FEC.Data[936] := 273.18;
   Prof_FEC.Data[937] := 251.28;
   Prof_FEC.Data[938] := 235.91;
   Prof_FEC.Data[939] := 224.8;
   Prof_FEC.Data[940] := 41.084;
   Prof_FEC.Data[941] := 40.079;
   Prof_FEC.Data[942] := 38.801;
   Prof_FEC.Data[943] := 37.72;
   Prof_FEC.Data[944] := 38.026;
   Prof_FEC.Data[945] := 36.96;
   Prof_FEC.Data[946] := 37.986;
   Prof_FEC.Data[947] := 35.946;
   Prof_FEC.Data[948] := 40.907;
   Prof_FEC.Data[949] := 41.802;
   Prof_FEC.Data[950] := 41.211;
   Prof_FEC.Data[951] := 40.913;
   Prof_FEC.Data[952] := 41.099;
   Prof_FEC.Data[953] := 38.1;
   Prof_FEC.Data[954] := 39.037;
   Prof_FEC.Data[955] := 38.068;
   Prof_FEC.Data[956] := 41.886;
   Prof_FEC.Data[957] := 41.446;
   Prof_FEC.Data[958] := 42.211;
   Prof_FEC.Data[959] := 41.845;
   Prof_FEC.Data[960] := 41.54;
   Prof_FEC.Data[961] := 42.515;
   Prof_FEC.Data[962] := 40.592;
   Prof_FEC.Data[963] := 43.014;
   Prof_FEC.Data[964] := 42.632;
   Prof_FEC.Data[965] := 41.208;
   Prof_FEC.Data[966] := 41.964;
   Prof_FEC.Data[967] := 40.41;
   Prof_FEC.Data[968] := 41.73;
   Prof_FEC.Data[969] := 42.281;
   Prof_FEC.Data[970] := 39.995;
   Prof_FEC.Data[971] := 39.995;
   Prof_FEC.Data[972] := 44.187;
   Prof_FEC.Data[973] := 47.132;
   Prof_FEC.Data[974] := 44.583;
   Prof_FEC.Data[975] := 44.8;
   Prof_FEC.Data[976] := 45.313;
   Prof_FEC.Data[977] := 41.308;
   Prof_FEC.Data[978] := 40.704;
   Prof_FEC.Data[979] := 41.699;
   Prof_FEC.Data[980] := 267.76;
   Prof_FEC.Data[981] := 317.35;
   Prof_FEC.Data[982] := 288.51;
   Prof_FEC.Data[983] := 273.95;
   Prof_FEC.Data[984] := 278.64;
   Prof_FEC.Data[985] := 218.73;
   Prof_FEC.Data[986] := 267.79;
   Prof_FEC.Data[987] := 273.85;
   Prof_FEC.Data[988] := 341.92;
   Prof_FEC.Data[989] := 353.15;
   Prof_FEC.Data[990] := 382.56;
   Prof_FEC.Data[991] := 372.59;
   Prof_FEC.Data[992] := 292.38;
   Prof_FEC.Data[993] := 287.67;
   Prof_FEC.Data[994] := 231.66;
   Prof_FEC.Data[995] := 282.21;
   Prof_FEC.Data[996] := 311.99;
   Prof_FEC.Data[997] := 338.5;
   Prof_FEC.Data[998] := 341.54;
   Prof_FEC.Data[999] := 313.02;
   Prof_FEC.Data[1000] := 303.97;
   Prof_FEC.Data[1001] := 341.66;
   Prof_FEC.Data[1002] := 314.71;
   Prof_FEC.Data[1003] := 359.5;
   Prof_FEC.Data[1004] := 340.78;
   Prof_FEC.Data[1005] := 373.27;
   Prof_FEC.Data[1006] := 353.28;
   Prof_FEC.Data[1007] := 327.86;
   Prof_FEC.Data[1008] := 289.59;
   Prof_FEC.Data[1009] := 263.97;
   Prof_FEC.Data[1010] := 254.34;
   Prof_FEC.Data[1011] := 286.36;
   Prof_FEC.Data[1012] := 249.6;
   Prof_FEC.Data[1013] := 241.63;
   Prof_FEC.Data[1014] := 282.42;
   Prof_FEC.Data[1015] := 302.78;
   Prof_FEC.Data[1016] := 305.85;
   Prof_FEC.Data[1017] := 268.56;
   Prof_FEC.Data[1018] := 249.07;
   Prof_FEC.Data[1019] := 250.66;
   Prof_FEC.Data[1020] := 267.91;
   Prof_FEC.Data[1021] := 274.46;
   Prof_FEC.Data[1022] := 260.83;
   Prof_FEC.Data[1023] := 253.06;
   Prof_FEC.Data[1024] := 220.9;
   Prof_FEC.Data[1025] := 211.49;
   Prof_FEC.Data[1026] := 221.01;
   Prof_FEC.Data[1027] := 226.58;
   Prof_FEC.Data[1028] := 273.65;
   Prof_FEC.Data[1029] := 286.2;
   Prof_FEC.Data[1030] := 273.19;
   Prof_FEC.Data[1031] := 275.69;
   Prof_FEC.Data[1032] := 310.43;
   Prof_FEC.Data[1033] := 288.34;
   Prof_FEC.Data[1034] := 332.78;
   Prof_FEC.Data[1035] := 311.66;
   Prof_FEC.Data[1036] := 44.076;
   Prof_FEC.Data[1037] := 46.338;
   Prof_FEC.Data[1038] := 44.021;
   Prof_FEC.Data[1039] := 46.373;
   Prof_FEC.Data[1040] := 45.752;
   Prof_FEC.Data[1041] := 50.0;
   Prof_FEC.Data[1042] := 50.0;
   Prof_FEC.Data[1043] := 46.194;
   Prof_FEC.Data[1044] := 44.029;
   Prof_FEC.Data[1045] := 45.361;
   Prof_FEC.Data[1046] := 42.191;
   Prof_FEC.Data[1047] := 44.109;
   Prof_FEC.Data[1048] := 43.526;
   Prof_FEC.Data[1049] := 44.218;
   Prof_FEC.Data[1050] := 44.652;
   Prof_FEC.Data[1051] := 43.306;
   Prof_FEC.Data[1052] := 41.161;
   Prof_FEC.Data[1053] := 36.829;
   Prof_FEC.Data[1054] := 41.06;
   Prof_FEC.Data[1055] := 39.562;
   Prof_FEC.Data[1056] := 45.987;
   Prof_FEC.Data[1057] := 42.254;
   Prof_FEC.Data[1058] := 46.048;
   Prof_FEC.Data[1059] := 45.769;
   Prof_FEC.Data[1060] := 43.262;
   Prof_FEC.Data[1061] := 43.505;
   Prof_FEC.Data[1062] := 44.086;
   Prof_FEC.Data[1063] := 44.927;
   Prof_FEC.Data[1064] := 46.993;
   Prof_FEC.Data[1065] := 50.0;
   Prof_FEC.Data[1066] := 50.0;
   Prof_FEC.Data[1067] := 50.0;
   Prof_FEC.Data[1068] := 48.38;
   Prof_FEC.Data[1069] := 46.334;
   Prof_FEC.Data[1070] := 45.352;
   Prof_FEC.Data[1071] := 50.0;
   Prof_FEC.Data[1072] := 50.0;
   Prof_FEC.Data[1073] := 50.0;
   Prof_FEC.Data[1074] := 50.0;
   Prof_FEC.Data[1075] := 50.0;
   Prof_FEC.Data[1076] := 343.88;
   Prof_FEC.Data[1077] := 276.6;
   Prof_FEC.Data[1078] := 277.09;
   Prof_FEC.Data[1079] := 306.26;
   Prof_FEC.Data[1080] := 282.63;
   Prof_FEC.Data[1081] := 319.68;
   Prof_FEC.Data[1082] := 331.81;
   Prof_FEC.Data[1083] := 293.38;
   Prof_FEC.Data[1084] := 264.96;
   Prof_FEC.Data[1085] := 269.32;
   Prof_FEC.Data[1086] := 261.4;
   Prof_FEC.Data[1087] := 237.31;
   Prof_FEC.Data[1088] := 237.03;
   Prof_FEC.Data[1089] := 202.12;
   Prof_FEC.Data[1090] := 187.81;
   Prof_FEC.Data[1091] := 202.7;
   Prof_FEC.Data[1092] := 170.03;
   Prof_FEC.Data[1093] := 149.46;
   Prof_FEC.Data[1094] := 171.4;
   Prof_FEC.Data[1095] := 191.13;
   Prof_FEC.Data[1096] := 221.65;
   Prof_FEC.Data[1097] := 239.58;
   Prof_FEC.Data[1098] := 220.51;
   Prof_FEC.Data[1099] := 209.37;
   Prof_FEC.Data[1100] := 168.01;
   Prof_FEC.Data[1101] := 167.58;
   Prof_FEC.Data[1102] := 161.67;
   Prof_FEC.Data[1103] := 170.39;
   Prof_FEC.Data[1104] := 185.36;
   Prof_FEC.Data[1105] := 235.04;
   Prof_FEC.Data[1106] := 169.17;
   Prof_FEC.Data[1107] := 185.62;
   Prof_FEC.Data[1108] := 154.96;
   Prof_FEC.Data[1109] := 158.08;
   Prof_FEC.Data[1110] := 146.87;
   Prof_FEC.Data[1111] := 155.1;
   Prof_FEC.Data[1112] := 195.69;
   Prof_FEC.Data[1113] := 206.16;
   Prof_FEC.Data[1114] := 198.86;
   Prof_FEC.Data[1115] := 198.48;
   Prof_FEC.Data[1116] := 158.56;
   Prof_FEC.Data[1117] := 157.48;
   Prof_FEC.Data[1118] := 174.9;
   Prof_FEC.Data[1119] := 185.12;
   Prof_FEC.Data[1120] := 261.63;
   Prof_FEC.Data[1121] := 257.58;
   Prof_FEC.Data[1122] := 272.92;
   Prof_FEC.Data[1123] := 276.31;
   Prof_FEC.Data[1124] := 302.74;
   Prof_FEC.Data[1125] := 293.63;
   Prof_FEC.Data[1126] := 276.29;
   Prof_FEC.Data[1127] := 315.21;
   Prof_FEC.Data[1128] := 307.15;
   Prof_FEC.Data[1129] := 344.1;
   Prof_FEC.Data[1130] := 348.66;
   Prof_FEC.Data[1131] := 352.85;
   Prof_FEC.Data[1132] := 45.874;
   Prof_FEC.Data[1133] := 48.345;
   Prof_FEC.Data[1134] := 46.881;
   Prof_FEC.Data[1135] := 48.553;
   Prof_FEC.Data[1136] := 46.393;
   Prof_FEC.Data[1137] := 47.929;
   Prof_FEC.Data[1138] := 50.0;
   Prof_FEC.Data[1139] := 50.0;
   Prof_FEC.Data[1140] := 48.298;
   Prof_FEC.Data[1141] := 50.0;
   Prof_FEC.Data[1142] := 47.419;
   Prof_FEC.Data[1143] := 48.943;
   Prof_FEC.Data[1144] := 50.0;
   Prof_FEC.Data[1145] := 50.0;
   Prof_FEC.Data[1146] := 50.0;
   Prof_FEC.Data[1147] := 50.0;
   Prof_FEC.Data[1148] := 50.0;
   Prof_FEC.Data[1149] := 47.395;
   Prof_FEC.Data[1150] := 47.988;
   Prof_FEC.Data[1151] := 50.0;
   Prof_FEC.Data[1152] := 50.0;
   Prof_FEC.Data[1153] := 50.0;
   Prof_FEC.Data[1154] := 50.0;
   Prof_FEC.Data[1155] := 50.0;
   Prof_FEC.Data[1156] := 50.0;
   Prof_FEC.Data[1157] := 49.565;
   Prof_FEC.Data[1158] := 50.0;
   Prof_FEC.Data[1159] := 50.0;
   Prof_FEC.Data[1160] := 50.0;
   Prof_FEC.Data[1161] := 50.0;
   Prof_FEC.Data[1162] := 50.0;
   Prof_FEC.Data[1163] := 50.0;
   Prof_FEC.Data[1164] := 49.623;
   Prof_FEC.Data[1165] := 47.95;
   Prof_FEC.Data[1166] := 49.51;
   Prof_FEC.Data[1167] := 50.0;
   Prof_FEC.Data[1168] := 50.0;
   Prof_FEC.Data[1169] := 50.0;
   Prof_FEC.Data[1170] := 50.0;
   Prof_FEC.Data[1171] := 50.0;
   Prof_FEC.Data[1172] := 346.66;
   Prof_FEC.Data[1173] := 335.08;
   Prof_FEC.Data[1174] := 333.85;
   Prof_FEC.Data[1175] := 308.36;
   Prof_FEC.Data[1176] := 379.12;
   Prof_FEC.Data[1177] := 418.58;
   Prof_FEC.Data[1178] := 370.95;
   Prof_FEC.Data[1179] := 437.4;
   Prof_FEC.Data[1180] := 467.47;
   Prof_FEC.Data[1181] := 536.25;
   Prof_FEC.Data[1182] := 552.01;
   Prof_FEC.Data[1183] := 577.38;
   Prof_FEC.Data[1184] := 553.14;
   Prof_FEC.Data[1185] := 564.29;
   Prof_FEC.Data[1186] := 600.41;
   Prof_FEC.Data[1187] := 638.88;
   Prof_FEC.Data[1188] := 643.54;
   Prof_FEC.Data[1189] := 718.29;
   Prof_FEC.Data[1190] := 674.3;
   Prof_FEC.Data[1191] := 677.75;
   Prof_FEC.Data[1192] := 664.48;
   Prof_FEC.Data[1193] := 636.75;
   Prof_FEC.Data[1194] := 680.46;
   Prof_FEC.Data[1195] := 644.66;
   Prof_FEC.Data[1196] := 666.58;
   Prof_FEC.Data[1197] := 691.69;
   Prof_FEC.Data[1198] := 619.25;
   Prof_FEC.Data[1199] := 657.49;
   Prof_FEC.Data[1200] := 639.27;
   Prof_FEC.Data[1201] := 631.76;
   Prof_FEC.Data[1202] := 590.65;
   Prof_FEC.Data[1203] := 556.39;
   Prof_FEC.Data[1204] := 584.07;
   Prof_FEC.Data[1205] := 598.69;
   Prof_FEC.Data[1206] := 655.75;
   Prof_FEC.Data[1207] := 616.22;
   Prof_FEC.Data[1208] := 557.33;
   Prof_FEC.Data[1209] := 517.14;
   Prof_FEC.Data[1210] := 558.55;
   Prof_FEC.Data[1211] := 620.38;
   Prof_FEC.Data[1212] := 619.44;
   Prof_FEC.Data[1213] := 574.65;
   Prof_FEC.Data[1214] := 680.51;
   Prof_FEC.Data[1215] := 635.81;
   Prof_FEC.Data[1216] := 587.69;
   Prof_FEC.Data[1217] := 637.69;
   Prof_FEC.Data[1218] := 650.52;
   Prof_FEC.Data[1219] := 556.97;
   Prof_FEC.Data[1220] := 428.74;
   Prof_FEC.Data[1221] := 391.72;
   Prof_FEC.Data[1222] := 357.99;
   Prof_FEC.Data[1223] := 347.31;
   Prof_FEC.Data[1224] := 349.11;
   Prof_FEC.Data[1225] := 321.45;
   Prof_FEC.Data[1226] := 324.29;
   Prof_FEC.Data[1227] := 293.91;
   Prof_FEC.Data[1228] := 49.81;
   Prof_FEC.Data[1229] := 50.0;
   Prof_FEC.Data[1230] := 50.0;
   Prof_FEC.Data[1231] := 50.0;
   Prof_FEC.Data[1232] := 48.891;
   Prof_FEC.Data[1233] := 50.0;
   Prof_FEC.Data[1234] := 48.222;
   Prof_FEC.Data[1235] := 48.49;
   Prof_FEC.Data[1236] := 50.0;
   Prof_FEC.Data[1237] := 50.0;
   Prof_FEC.Data[1238] := 50.0;
   Prof_FEC.Data[1239] := 50.0;
   Prof_FEC.Data[1240] := 46.469;
   Prof_FEC.Data[1241] := 47.92;
   Prof_FEC.Data[1242] := 45.351;
   Prof_FEC.Data[1243] := 46.449;
   Prof_FEC.Data[1244] := 49.791;
   Prof_FEC.Data[1245] := 50.0;
   Prof_FEC.Data[1246] := 47.006;
   Prof_FEC.Data[1247] := 49.828;
   Prof_FEC.Data[1248] := 41.868;
   Prof_FEC.Data[1249] := 44.705;
   Prof_FEC.Data[1250] := 41.45;
   Prof_FEC.Data[1251] := 42.297;
   Prof_FEC.Data[1252] := 45.338;
   Prof_FEC.Data[1253] := 45.547;
   Prof_FEC.Data[1254] := 42.009;
   Prof_FEC.Data[1255] := 45.826;
   Prof_FEC.Data[1256] := 44.373;
   Prof_FEC.Data[1257] := 42.367;
   Prof_FEC.Data[1258] := 40.681;
   Prof_FEC.Data[1259] := 39.686;
   Prof_FEC.Data[1260] := 40.095;
   Prof_FEC.Data[1261] := 40.725;
   Prof_FEC.Data[1262] := 45.116;
   Prof_FEC.Data[1263] := 44.975;
   Prof_FEC.Data[1264] := 42.353;
   Prof_FEC.Data[1265] := 42.292;
   Prof_FEC.Data[1266] := 41.993;
   Prof_FEC.Data[1267] := 41.815;
   Prof_FEC.Data[1268] := 245.69;
   Prof_FEC.Data[1269] := 274.47;
   Prof_FEC.Data[1270] := 294.63;
   Prof_FEC.Data[1271] := 310.82;
   Prof_FEC.Data[1272] := 330.41;
   Prof_FEC.Data[1273] := 341.4;
   Prof_FEC.Data[1274] := 279.25;
   Prof_FEC.Data[1275] := 347.41;
   Prof_FEC.Data[1276] := 387.2;
   Prof_FEC.Data[1277] := 461.69;
   Prof_FEC.Data[1278] := 411.45;
   Prof_FEC.Data[1279] := 402.32;
   Prof_FEC.Data[1280] := 496.79;
   Prof_FEC.Data[1281] := 500.77;
   Prof_FEC.Data[1282] := 450.71;
   Prof_FEC.Data[1283] := 493.87;
   Prof_FEC.Data[1284] := 592.78;
   Prof_FEC.Data[1285] := 536.33;
   Prof_FEC.Data[1286] := 588.07;
   Prof_FEC.Data[1287] := 641.5;
   Prof_FEC.Data[1288] := 558.41;
   Prof_FEC.Data[1289] := 633.34;
   Prof_FEC.Data[1290] := 592.09;
   Prof_FEC.Data[1291] := 616.68;
   Prof_FEC.Data[1292] := 605.73;
   Prof_FEC.Data[1293] := 618.94;
   Prof_FEC.Data[1294] := 616.0;
   Prof_FEC.Data[1295] := 642.12;
   Prof_FEC.Data[1296] := 656.39;
   Prof_FEC.Data[1297] := 570.61;
   Prof_FEC.Data[1298] := 576.67;
   Prof_FEC.Data[1299] := 609.67;
   Prof_FEC.Data[1300] := 648.23;
   Prof_FEC.Data[1301] := 714.64;
   Prof_FEC.Data[1302] := 714.68;
   Prof_FEC.Data[1303] := 703.72;
   Prof_FEC.Data[1304] := 641.36;
   Prof_FEC.Data[1305] := 637.64;
   Prof_FEC.Data[1306] := 669.93;
   Prof_FEC.Data[1307] := 639.96;
   Prof_FEC.Data[1308] := 571.97;
   Prof_FEC.Data[1309] := 673.36;
   Prof_FEC.Data[1310] := 649.85;
   Prof_FEC.Data[1311] := 738.51;
   Prof_FEC.Data[1312] := 807.53;
   Prof_FEC.Data[1313] := 700.68;
   Prof_FEC.Data[1314] := 774.95;
   Prof_FEC.Data[1315] := 667.65;
   Prof_FEC.Data[1316] := 458.36;
   Prof_FEC.Data[1317] := 438.58;
   Prof_FEC.Data[1318] := 340.71;
   Prof_FEC.Data[1319] := 351.08;
   Prof_FEC.Data[1320] := 286.57;
   Prof_FEC.Data[1321] := 245.11;
   Prof_FEC.Data[1322] := 281.93;
   Prof_FEC.Data[1323] := 247.85;
   Prof_FEC.Data[1324] := 43.541;
   Prof_FEC.Data[1325] := 44.758;
   Prof_FEC.Data[1326] := 45.046;
   Prof_FEC.Data[1327] := 46.627;
   Prof_FEC.Data[1328] := 44.031;
   Prof_FEC.Data[1329] := 44.011;
   Prof_FEC.Data[1330] := 43.231;
   Prof_FEC.Data[1331] := 38.834;
   Prof_FEC.Data[1332] := 43.238;
   Prof_FEC.Data[1333] := 40.282;
   Prof_FEC.Data[1334] := 37.897;
   Prof_FEC.Data[1335] := 41.441;
   Prof_FEC.Data[1336] := 38.746;
   Prof_FEC.Data[1337] := 37.925;
   Prof_FEC.Data[1338] := 37.576;
   Prof_FEC.Data[1339] := 37.523;
   Prof_FEC.Data[1340] := 39.74;
   Prof_FEC.Data[1341] := 41.639;
   Prof_FEC.Data[1342] := 40.508;
   Prof_FEC.Data[1343] := 39.558;
   Prof_FEC.Data[1344] := 40.986;
   Prof_FEC.Data[1345] := 41.139;
   Prof_FEC.Data[1346] := 39.577;
   Prof_FEC.Data[1347] := 39.532;
   Prof_FEC.Data[1348] := 40.801;
   Prof_FEC.Data[1349] := 39.649;
   Prof_FEC.Data[1350] := 41.681;
   Prof_FEC.Data[1351] := 39.168;
   Prof_FEC.Data[1352] := 37.814;
   Prof_FEC.Data[1353] := 35.978;
   Prof_FEC.Data[1354] := 37.618;
   Prof_FEC.Data[1355] := 37.61;
   Prof_FEC.Data[1356] := 38.979;
   Prof_FEC.Data[1357] := 41.857;
   Prof_FEC.Data[1358] := 40.187;
   Prof_FEC.Data[1359] := 37.132;
   Prof_FEC.Data[1360] := 39.955;
   Prof_FEC.Data[1361] := 36.961;
   Prof_FEC.Data[1362] := 38.953;
   Prof_FEC.Data[1363] := 38.771;
   Prof_FEC.Data[1364] := 248.93;
   Prof_FEC.Data[1365] := 243.32;
   Prof_FEC.Data[1366] := 262.85;
   Prof_FEC.Data[1367] := 304.98;
   Prof_FEC.Data[1368] := 349.72;
   Prof_FEC.Data[1369] := 423.12;
   Prof_FEC.Data[1370] := 405.04;
   Prof_FEC.Data[1371] := 443.58;
   Prof_FEC.Data[1372] := 460.14;
   Prof_FEC.Data[1373] := 513.79;
   Prof_FEC.Data[1374] := 513.42;
   Prof_FEC.Data[1375] := 610.74;
   Prof_FEC.Data[1376] := 559.36;
   Prof_FEC.Data[1377] := 606.73;
   Prof_FEC.Data[1378] := 592.74;
   Prof_FEC.Data[1379] := 676.69;
   Prof_FEC.Data[1380] := 700.62;
   Prof_FEC.Data[1381] := 756.2;
   Prof_FEC.Data[1382] := 709.31;
   Prof_FEC.Data[1383] := 770.89;
   Prof_FEC.Data[1384] := 752.41;
   Prof_FEC.Data[1385] := 719.2;
   Prof_FEC.Data[1386] := 700.3;
   Prof_FEC.Data[1387] := 713.47;
   Prof_FEC.Data[1388] := 681.02;
   Prof_FEC.Data[1389] := 678.77;
   Prof_FEC.Data[1390] := 735.62;
   Prof_FEC.Data[1391] := 680.6;
   Prof_FEC.Data[1392] := 685.99;
   Prof_FEC.Data[1393] := 709.12;
   Prof_FEC.Data[1394] := 620.42;
   Prof_FEC.Data[1395] := 653.23;
   Prof_FEC.Data[1396] := 678.39;
   Prof_FEC.Data[1397] := 665.12;
   Prof_FEC.Data[1398] := 667.9;
   Prof_FEC.Data[1399] := 626.61;
   Prof_FEC.Data[1400] := 694.11;
   Prof_FEC.Data[1401] := 636.51;
   Prof_FEC.Data[1402] := 644.14;
   Prof_FEC.Data[1403] := 633.12;
   Prof_FEC.Data[1404] := 668.63;
   Prof_FEC.Data[1405] := 636.63;
   Prof_FEC.Data[1406] := 638.53;
   Prof_FEC.Data[1407] := 717.97;
   Prof_FEC.Data[1408] := 707.55;
   Prof_FEC.Data[1409] := 728.57;
   Prof_FEC.Data[1410] := 676.85;
   Prof_FEC.Data[1411] := 579.31;
   Prof_FEC.Data[1412] := 443.58;
   Prof_FEC.Data[1413] := 387.07;
   Prof_FEC.Data[1414] := 385.49;
   Prof_FEC.Data[1415] := 334.02;
   Prof_FEC.Data[1416] := 302.04;
   Prof_FEC.Data[1417] := 283.71;
   Prof_FEC.Data[1418] := 269.28;
   Prof_FEC.Data[1419] := 288.69;
   Prof_FEC.Data[1420] := 47.17;
   Prof_FEC.Data[1421] := 49.817;
   Prof_FEC.Data[1422] := 48.096;
   Prof_FEC.Data[1423] := 48.799;
   Prof_FEC.Data[1424] := 44.355;
   Prof_FEC.Data[1425] := 47.509;
   Prof_FEC.Data[1426] := 44.71;
   Prof_FEC.Data[1427] := 45.721;
   Prof_FEC.Data[1428] := 48.192;
   Prof_FEC.Data[1429] := 47.619;
   Prof_FEC.Data[1430] := 48.057;
   Prof_FEC.Data[1431] := 49.208;
   Prof_FEC.Data[1432] := 44.057;
   Prof_FEC.Data[1433] := 43.768;
   Prof_FEC.Data[1434] := 42.188;
   Prof_FEC.Data[1435] := 42.575;
   Prof_FEC.Data[1436] := 46.265;
   Prof_FEC.Data[1437] := 49.647;
   Prof_FEC.Data[1438] := 50.0;
   Prof_FEC.Data[1439] := 47.289;
   Prof_FEC.Data[1440] := 48.223;
   Prof_FEC.Data[1441] := 45.332;
   Prof_FEC.Data[1442] := 45.785;
   Prof_FEC.Data[1443] := 45.275;
   Prof_FEC.Data[1444] := 50.0;
   Prof_FEC.Data[1445] := 50.0;
   Prof_FEC.Data[1446] := 50.0;
   Prof_FEC.Data[1447] := 50.0;
   Prof_FEC.Data[1448] := 46.883;
   Prof_FEC.Data[1449] := 43.314;
   Prof_FEC.Data[1450] := 48.246;
   Prof_FEC.Data[1451] := 44.93;
   Prof_FEC.Data[1452] := 50.0;
   Prof_FEC.Data[1453] := 50.0;
   Prof_FEC.Data[1454] := 50.0;
   Prof_FEC.Data[1455] := 48.26;
   Prof_FEC.Data[1456] := 44.769;
   Prof_FEC.Data[1457] := 44.43;
   Prof_FEC.Data[1458] := 41.078;
   Prof_FEC.Data[1459] := 43.537;
   Prof_FEC.Data[1460] := 331.56;
   Prof_FEC.Data[1461] := 384.93;
   Prof_FEC.Data[1462] := 348.44;
   Prof_FEC.Data[1463] := 385.17;
   Prof_FEC.Data[1464] := 414.66;
   Prof_FEC.Data[1465] := 381.47;
   Prof_FEC.Data[1466] := 476.75;
   Prof_FEC.Data[1467] := 459.41;
   Prof_FEC.Data[1468] := 526.59;
   Prof_FEC.Data[1469] := 570.48;
   Prof_FEC.Data[1470] := 561.18;
   Prof_FEC.Data[1471] := 515.0;
   Prof_FEC.Data[1472] := 595.45;
   Prof_FEC.Data[1473] := 480.3;
   Prof_FEC.Data[1474] := 525.31;
   Prof_FEC.Data[1475] := 560.33;
   Prof_FEC.Data[1476] := 601.83;
   Prof_FEC.Data[1477] := 696.95;
   Prof_FEC.Data[1478] := 598.31;
   Prof_FEC.Data[1479] := 732.39;
   Prof_FEC.Data[1480] := 692.09;
   Prof_FEC.Data[1481] := 663.17;
   Prof_FEC.Data[1482] := 654.84;
   Prof_FEC.Data[1483] := 737.02;
   Prof_FEC.Data[1484] := 743.97;
   Prof_FEC.Data[1485] := 779.49;
   Prof_FEC.Data[1486] := 753.67;
   Prof_FEC.Data[1487] := 787.23;
   Prof_FEC.Data[1488] := 687.99;
   Prof_FEC.Data[1489] := 673.92;
   Prof_FEC.Data[1490] := 683.87;
   Prof_FEC.Data[1491] := 654.51;
   Prof_FEC.Data[1492] := 726.98;
   Prof_FEC.Data[1493] := 765.27;
   Prof_FEC.Data[1494] := 749.55;
   Prof_FEC.Data[1495] := 747.21;
   Prof_FEC.Data[1496] := 736.7;
   Prof_FEC.Data[1497] := 619.37;
   Prof_FEC.Data[1498] := 695.2;
   Prof_FEC.Data[1499] := 689.46;
   Prof_FEC.Data[1500] := 720.94;
   Prof_FEC.Data[1501] := 670.68;
   Prof_FEC.Data[1502] := 744.18;
   Prof_FEC.Data[1503] := 674.61;
   Prof_FEC.Data[1504] := 768.02;
   Prof_FEC.Data[1505] := 773.92;
   Prof_FEC.Data[1506] := 785.39;
   Prof_FEC.Data[1507] := 576.63;
   Prof_FEC.Data[1508] := 518.95;
   Prof_FEC.Data[1509] := 423.4;
   Prof_FEC.Data[1510] := 350.57;
   Prof_FEC.Data[1511] := 344.44;
   Prof_FEC.Data[1512] := 297.4;
   Prof_FEC.Data[1513] := 270.07;
   Prof_FEC.Data[1514] := 243.69;
   Prof_FEC.Data[1515] := 264.76;
   Prof_FEC.Data[1516] := 39.313;
   Prof_FEC.Data[1517] := 43.751;
   Prof_FEC.Data[1518] := 40.956;
   Prof_FEC.Data[1519] := 43.177;
   Prof_FEC.Data[1520] := 44.765;
   Prof_FEC.Data[1521] := 41.81;
   Prof_FEC.Data[1522] := 42.317;
   Prof_FEC.Data[1523] := 42.331;
   Prof_FEC.Data[1524] := 45.655;
   Prof_FEC.Data[1525] := 42.807;
   Prof_FEC.Data[1526] := 40.799;
   Prof_FEC.Data[1527] := 40.101;
   Prof_FEC.Data[1528] := 35.822;
   Prof_FEC.Data[1529] := 39.236;
   Prof_FEC.Data[1530] := 40.036;
   Prof_FEC.Data[1531] := 39.258;
   Prof_FEC.Data[1532] := 42.501;
   Prof_FEC.Data[1533] := 44.856;
   Prof_FEC.Data[1534] := 45.402;
   Prof_FEC.Data[1535] := 42.666;
   Prof_FEC.Data[1536] := 41.427;
   Prof_FEC.Data[1537] := 42.113;
   Prof_FEC.Data[1538] := 42.326;
   Prof_FEC.Data[1539] := 43.826;
   Prof_FEC.Data[1540] := 45.613;
   Prof_FEC.Data[1541] := 48.888;
   Prof_FEC.Data[1542] := 42.941;
   Prof_FEC.Data[1543] := 43.606;
   Prof_FEC.Data[1544] := 37.865;
   Prof_FEC.Data[1545] := 41.188;
   Prof_FEC.Data[1546] := 38.783;
   Prof_FEC.Data[1547] := 38.378;
   Prof_FEC.Data[1548] := 39.922;
   Prof_FEC.Data[1549] := 36.865;
   Prof_FEC.Data[1550] := 39.602;
   Prof_FEC.Data[1551] := 42.225;
   Prof_FEC.Data[1552] := 40.479;
   Prof_FEC.Data[1553] := 41.718;
   Prof_FEC.Data[1554] := 37.268;
   Prof_FEC.Data[1555] := 39.389;
   Prof_FEC.Data[1556] := 217.2;
   Prof_FEC.Data[1557] := 215.66;
   Prof_FEC.Data[1558] := 235.16;
   Prof_FEC.Data[1559] := 248.61;
   Prof_FEC.Data[1560] := 300.01;
   Prof_FEC.Data[1561] := 318.85;
   Prof_FEC.Data[1562] := 335.06;
   Prof_FEC.Data[1563] := 397.96;
   Prof_FEC.Data[1564] := 437.56;
   Prof_FEC.Data[1565] := 438.1;
   Prof_FEC.Data[1566] := 501.62;
   Prof_FEC.Data[1567] := 544.11;
   Prof_FEC.Data[1568] := 548.93;
   Prof_FEC.Data[1569] := 505.75;
   Prof_FEC.Data[1570] := 457.03;
   Prof_FEC.Data[1571] := 559.36;
   Prof_FEC.Data[1572] := 620.63;
   Prof_FEC.Data[1573] := 587.33;
   Prof_FEC.Data[1574] := 653.36;
   Prof_FEC.Data[1575] := 693.94;
   Prof_FEC.Data[1576] := 719.77;
   Prof_FEC.Data[1577] := 667.78;
   Prof_FEC.Data[1578] := 743.75;
   Prof_FEC.Data[1579] := 760.63;
   Prof_FEC.Data[1580] := 730.56;
   Prof_FEC.Data[1581] := 743.92;
   Prof_FEC.Data[1582] := 693.92;
   Prof_FEC.Data[1583] := 689.24;
   Prof_FEC.Data[1584] := 623.36;
   Prof_FEC.Data[1585] := 555.63;
   Prof_FEC.Data[1586] := 646.63;
   Prof_FEC.Data[1587] := 644.12;
   Prof_FEC.Data[1588] := 635.72;
   Prof_FEC.Data[1589] := 624.64;
   Prof_FEC.Data[1590] := 626.05;
   Prof_FEC.Data[1591] := 634.16;
   Prof_FEC.Data[1592] := 658.13;
   Prof_FEC.Data[1593] := 640.64;
   Prof_FEC.Data[1594] := 663.39;
   Prof_FEC.Data[1595] := 668.04;
   Prof_FEC.Data[1596] := 625.8;
   Prof_FEC.Data[1597] := 651.86;
   Prof_FEC.Data[1598] := 568.48;
   Prof_FEC.Data[1599] := 552.16;
   Prof_FEC.Data[1600] := 740.52;
   Prof_FEC.Data[1601] := 665.07;
   Prof_FEC.Data[1602] := 548.25;
   Prof_FEC.Data[1603] := 529.77;
   Prof_FEC.Data[1604] := 377.7;
   Prof_FEC.Data[1605] := 301.4;
   Prof_FEC.Data[1606] := 264.49;
   Prof_FEC.Data[1607] := 243.83;
   Prof_FEC.Data[1608] := 241.44;
   Prof_FEC.Data[1609] := 222.71;
   Prof_FEC.Data[1610] := 222.38;
   Prof_FEC.Data[1611] := 210.89;
   Prof_FEC.Data[1612] := 41.774;
   Prof_FEC.Data[1613] := 40.189;
   Prof_FEC.Data[1614] := 42.587;
   Prof_FEC.Data[1615] := 38.47;
   Prof_FEC.Data[1616] := 35.747;
   Prof_FEC.Data[1617] := 39.624;
   Prof_FEC.Data[1618] := 38.639;
   Prof_FEC.Data[1619] := 38.625;
   Prof_FEC.Data[1620] := 39.23;
   Prof_FEC.Data[1621] := 39.834;
   Prof_FEC.Data[1622] := 40.701;
   Prof_FEC.Data[1623] := 42.798;
   Prof_FEC.Data[1624] := 41.881;
   Prof_FEC.Data[1625] := 38.443;
   Prof_FEC.Data[1626] := 44.201;
   Prof_FEC.Data[1627] := 41.771;
   Prof_FEC.Data[1628] := 46.58;
   Prof_FEC.Data[1629] := 44.587;
   Prof_FEC.Data[1630] := 45.351;
   Prof_FEC.Data[1631] := 44.285;
   Prof_FEC.Data[1632] := 42.278;
   Prof_FEC.Data[1633] := 39.23;
   Prof_FEC.Data[1634] := 41.167;
   Prof_FEC.Data[1635] := 43.32;
   Prof_FEC.Data[1636] := 43.432;
   Prof_FEC.Data[1637] := 43.034;
   Prof_FEC.Data[1638] := 43.137;
   Prof_FEC.Data[1639] := 42.443;
   Prof_FEC.Data[1640] := 42.008;
   Prof_FEC.Data[1641] := 43.467;
   Prof_FEC.Data[1642] := 44.079;
   Prof_FEC.Data[1643] := 42.055;
   Prof_FEC.Data[1644] := 48.538;
   Prof_FEC.Data[1645] := 46.533;
   Prof_FEC.Data[1646] := 48.241;
   Prof_FEC.Data[1647] := 44.681;
   Prof_FEC.Data[1648] := 43.223;
   Prof_FEC.Data[1649] := 44.315;
   Prof_FEC.Data[1650] := 41.095;
   Prof_FEC.Data[1651] := 43.459;
   Prof_FEC.Data[1652] := 314.37;
   Prof_FEC.Data[1653] := 303.72;
   Prof_FEC.Data[1654] := 305.29;
   Prof_FEC.Data[1655] := 348.37;
   Prof_FEC.Data[1656] := 331.65;
   Prof_FEC.Data[1657] := 293.46;
   Prof_FEC.Data[1658] := 299.95;
   Prof_FEC.Data[1659] := 305.67;
   Prof_FEC.Data[1660] := 414.37;
   Prof_FEC.Data[1661] := 430.71;
   Prof_FEC.Data[1662] := 466.04;
   Prof_FEC.Data[1663] := 421.51;
   Prof_FEC.Data[1664] := 353.7;
   Prof_FEC.Data[1665] := 306.55;
   Prof_FEC.Data[1666] := 284.95;
   Prof_FEC.Data[1667] := 305.79;
   Prof_FEC.Data[1668] := 366.59;
   Prof_FEC.Data[1669] := 357.83;
   Prof_FEC.Data[1670] := 360.0;
   Prof_FEC.Data[1671] := 392.56;
   Prof_FEC.Data[1672] := 382.91;
   Prof_FEC.Data[1673] := 382.11;
   Prof_FEC.Data[1674] := 407.14;
   Prof_FEC.Data[1675] := 396.69;
   Prof_FEC.Data[1676] := 362.19;
   Prof_FEC.Data[1677] := 374.45;
   Prof_FEC.Data[1678] := 357.09;
   Prof_FEC.Data[1679] := 355.92;
   Prof_FEC.Data[1680] := 287.07;
   Prof_FEC.Data[1681] := 269.62;
   Prof_FEC.Data[1682] := 220.37;
   Prof_FEC.Data[1683] := 227.0;
   Prof_FEC.Data[1684] := 261.66;
   Prof_FEC.Data[1685] := 272.23;
   Prof_FEC.Data[1686] := 249.62;
   Prof_FEC.Data[1687] := 244.34;
   Prof_FEC.Data[1688] := 256.03;
   Prof_FEC.Data[1689] := 221.83;
   Prof_FEC.Data[1690] := 247.05;
   Prof_FEC.Data[1691] := 245.21;
   Prof_FEC.Data[1692] := 247.55;
   Prof_FEC.Data[1693] := 231.56;
   Prof_FEC.Data[1694] := 234.89;
   Prof_FEC.Data[1695] := 191.04;
   Prof_FEC.Data[1696] := 169.13;
   Prof_FEC.Data[1697] := 162.61;
   Prof_FEC.Data[1698] := 157.02;
   Prof_FEC.Data[1699] := 186.3;
   Prof_FEC.Data[1700] := 218.08;
   Prof_FEC.Data[1701] := 242.93;
   Prof_FEC.Data[1702] := 235.85;
   Prof_FEC.Data[1703] := 249.02;
   Prof_FEC.Data[1704] := 255.77;
   Prof_FEC.Data[1705] := 227.69;
   Prof_FEC.Data[1706] := 237.15;
   Prof_FEC.Data[1707] := 213.09;
   Prof_FEC.Data[1708] := 38.285;
   Prof_FEC.Data[1709] := 38.585;
   Prof_FEC.Data[1710] := 40.036;
   Prof_FEC.Data[1711] := 38.163;
   Prof_FEC.Data[1712] := 38.293;
   Prof_FEC.Data[1713] := 40.463;
   Prof_FEC.Data[1714] := 36.484;
   Prof_FEC.Data[1715] := 37.325;
   Prof_FEC.Data[1716] := 34.758;
   Prof_FEC.Data[1717] := 37.891;
   Prof_FEC.Data[1718] := 37.618;
   Prof_FEC.Data[1719] := 39.685;
   Prof_FEC.Data[1720] := 40.379;
   Prof_FEC.Data[1721] := 41.635;
   Prof_FEC.Data[1722] := 45.444;
   Prof_FEC.Data[1723] := 41.835;
   Prof_FEC.Data[1724] := 41.948;
   Prof_FEC.Data[1725] := 40.107;
   Prof_FEC.Data[1726] := 39.252;
   Prof_FEC.Data[1727] := 42.538;
   Prof_FEC.Data[1728] := 43.187;
   Prof_FEC.Data[1729] := 43.07;
   Prof_FEC.Data[1730] := 43.112;
   Prof_FEC.Data[1731] := 42.238;
   Prof_FEC.Data[1732] := 40.756;
   Prof_FEC.Data[1733] := 40.258;
   Prof_FEC.Data[1734] := 41.165;
   Prof_FEC.Data[1735] := 43.805;
   Prof_FEC.Data[1736] := 41.15;
   Prof_FEC.Data[1737] := 43.529;
   Prof_FEC.Data[1738] := 44.109;
   Prof_FEC.Data[1739] := 41.298;
   Prof_FEC.Data[1740] := 41.453;
   Prof_FEC.Data[1741] := 40.338;
   Prof_FEC.Data[1742] := 41.795;
   Prof_FEC.Data[1743] := 42.058;
   Prof_FEC.Data[1744] := 41.748;
   Prof_FEC.Data[1745] := 43.955;
   Prof_FEC.Data[1746] := 40.794;
   Prof_FEC.Data[1747] := 42.64;
   Prof_FEC.Data[1748] := 244.32;
   Prof_FEC.Data[1749] := 254.73;
   Prof_FEC.Data[1750] := 247.34;
   Prof_FEC.Data[1751] := 256.6;
   Prof_FEC.Data[1752] := 264.29;
   Prof_FEC.Data[1753] := 279.93;
   Prof_FEC.Data[1754] := 278.29;
   Prof_FEC.Data[1755] := 275.43;
   Prof_FEC.Data[1756] := 257.49;
   Prof_FEC.Data[1757] := 228.72;
   Prof_FEC.Data[1758] := 218.18;
   Prof_FEC.Data[1759] := 193.68;
   Prof_FEC.Data[1760] := 160.39;
   Prof_FEC.Data[1761] := 155.78;
   Prof_FEC.Data[1762] := 127.38;
   Prof_FEC.Data[1763] := 133.79;
   Prof_FEC.Data[1764] := 133.42;
   Prof_FEC.Data[1765] := 108.95;
   Prof_FEC.Data[1766] := 106.76;
   Prof_FEC.Data[1767] := 116.01;
   Prof_FEC.Data[1768] := 108.36;
   Prof_FEC.Data[1769] := 137.08;
   Prof_FEC.Data[1770] := 127.71;
   Prof_FEC.Data[1771] := 118.36;
   Prof_FEC.Data[1772] := 117.67;
   Prof_FEC.Data[1773] := 102.75;
   Prof_FEC.Data[1774] := 104.67;
   Prof_FEC.Data[1775] := 106.73;
   Prof_FEC.Data[1776] := 119.04;
   Prof_FEC.Data[1777] := 130.37;
   Prof_FEC.Data[1778] := 111.31;
   Prof_FEC.Data[1779] := 124.02;
   Prof_FEC.Data[1780] := 98.34;
   Prof_FEC.Data[1781] := 113.9;
   Prof_FEC.Data[1782] := 105.94;
   Prof_FEC.Data[1783] := 106.98;
   Prof_FEC.Data[1784] := 122.42;
   Prof_FEC.Data[1785] := 119.33;
   Prof_FEC.Data[1786] := 118.03;
   Prof_FEC.Data[1787] := 122.2;
   Prof_FEC.Data[1788] := 102.51;
   Prof_FEC.Data[1789] := 94.45;
   Prof_FEC.Data[1790] := 109.68;
   Prof_FEC.Data[1791] := 130.15;
   Prof_FEC.Data[1792] := 159.58;
   Prof_FEC.Data[1793] := 173.58;
   Prof_FEC.Data[1794] := 197.97;
   Prof_FEC.Data[1795] := 228.33;
   Prof_FEC.Data[1796] := 223.68;
   Prof_FEC.Data[1797] := 238.19;
   Prof_FEC.Data[1798] := 267.8;
   Prof_FEC.Data[1799] := 273.29;
   Prof_FEC.Data[1800] := 268.08;
   Prof_FEC.Data[1801] := 283.23;
   Prof_FEC.Data[1802] := 325.44;
   Prof_FEC.Data[1803] := 287.06;
   Prof_FEC.Data[1804] := 40.4;
   Prof_FEC.Data[1805] := 40.478;
   Prof_FEC.Data[1806] := 40.205;
   Prof_FEC.Data[1807] := 42.619;
   Prof_FEC.Data[1808] := 43.622;
   Prof_FEC.Data[1809] := 41.93;
   Prof_FEC.Data[1810] := 45.305;
   Prof_FEC.Data[1811] := 43.209;
   Prof_FEC.Data[1812] := 41.556;
   Prof_FEC.Data[1813] := 40.547;
   Prof_FEC.Data[1814] := 40.422;
   Prof_FEC.Data[1815] := 39.503;
   Prof_FEC.Data[1816] := 41.029;
   Prof_FEC.Data[1817] := 39.23;
   Prof_FEC.Data[1818] := 41.379;
   Prof_FEC.Data[1819] := 39.293;
   Prof_FEC.Data[1820] := 39.504;
   Prof_FEC.Data[1821] := 36.708;
   Prof_FEC.Data[1822] := 36.181;
   Prof_FEC.Data[1823] := 37.796;
   Prof_FEC.Data[1824] := 39.781;
   Prof_FEC.Data[1825] := 37.202;
   Prof_FEC.Data[1826] := 38.329;
   Prof_FEC.Data[1827] := 38.739;
   Prof_FEC.Data[1828] := 38.461;
   Prof_FEC.Data[1829] := 37.362;
   Prof_FEC.Data[1830] := 40.23;
   Prof_FEC.Data[1831] := 38.853;
   Prof_FEC.Data[1832] := 39.902;
   Prof_FEC.Data[1833] := 40.227;
   Prof_FEC.Data[1834] := 40.502;
   Prof_FEC.Data[1835] := 40.606;
   Prof_FEC.Data[1836] := 38.466;
   Prof_FEC.Data[1837] := 37.51;
   Prof_FEC.Data[1838] := 38.87;
   Prof_FEC.Data[1839] := 37.859;
   Prof_FEC.Data[1840] := 42.166;
   Prof_FEC.Data[1841] := 42.681;
   Prof_FEC.Data[1842] := 44.4;
   Prof_FEC.Data[1843] := 43.613;
   Prof_FEC.Data[1844] := 294.01;
   Prof_FEC.Data[1845] := 269.82;
   Prof_FEC.Data[1846] := 260.38;
   Prof_FEC.Data[1847] := 261.77;
   Prof_FEC.Data[1848] := 284.95;
   Prof_FEC.Data[1849] := 277.73;
   Prof_FEC.Data[1850] := 266.54;
   Prof_FEC.Data[1851] := 267.19;
   Prof_FEC.Data[1852] := 224.86;
   Prof_FEC.Data[1853] := 190.26;
   Prof_FEC.Data[1854] := 199.84;
   Prof_FEC.Data[1855] := 187.43;
   Prof_FEC.Data[1856] := 144.18;
   Prof_FEC.Data[1857] := 102.79;
   Prof_FEC.Data[1858] := 111.4;
   Prof_FEC.Data[1859] := 102.16;
   Prof_FEC.Data[1860] := 107.39;
   Prof_FEC.Data[1861] := 106.93;
   Prof_FEC.Data[1862] := 88.62;
   Prof_FEC.Data[1863] := 109.44;
   Prof_FEC.Data[1864] := 117.67;
   Prof_FEC.Data[1865] := 135.62;
   Prof_FEC.Data[1866] := 127.74;
   Prof_FEC.Data[1867] := 117.95;
   Prof_FEC.Data[1868] := 120.15;
   Prof_FEC.Data[1869] := 94.06;
   Prof_FEC.Data[1870] := 111.86;
   Prof_FEC.Data[1871] := 100.72;
   Prof_FEC.Data[1872] := 116.22;
   Prof_FEC.Data[1873] := 121.43;
   Prof_FEC.Data[1874] := 125.75;
   Prof_FEC.Data[1875] := 129.51;
   Prof_FEC.Data[1876] := 94.66;
   Prof_FEC.Data[1877] := 99.86;
   Prof_FEC.Data[1878] := 108.31;
   Prof_FEC.Data[1879] := 94.02;
   Prof_FEC.Data[1880] := 105.07;
   Prof_FEC.Data[1881] := 110.06;
   Prof_FEC.Data[1882] := 117.6;
   Prof_FEC.Data[1883] := 109.74;
   Prof_FEC.Data[1884] := 89.51;
   Prof_FEC.Data[1885] := 83.69;
   Prof_FEC.Data[1886] := 104.66;
   Prof_FEC.Data[1887] := 107.5;
   Prof_FEC.Data[1888] := 120.19;
   Prof_FEC.Data[1889] := 139.2;
   Prof_FEC.Data[1890] := 149.83;
   Prof_FEC.Data[1891] := 185.36;
   Prof_FEC.Data[1892] := 195.46;
   Prof_FEC.Data[1893] := 244.18;
   Prof_FEC.Data[1894] := 254.08;
   Prof_FEC.Data[1895] := 250.03;
   Prof_FEC.Data[1896] := 224.36;
   Prof_FEC.Data[1897] := 229.18;
   Prof_FEC.Data[1898] := 223.71;
   Prof_FEC.Data[1899] := 252.92;
   Prof_FEC.Data[1900] := 36.389;
   Prof_FEC.Data[1901] := 36.914;
   Prof_FEC.Data[1902] := 37.863;
   Prof_FEC.Data[1903] := 35.113;
   Prof_FEC.Data[1904] := 37.029;
   Prof_FEC.Data[1905] := 34.587;
   Prof_FEC.Data[1906] := 39.12;
   Prof_FEC.Data[1907] := 34.629;
   Prof_FEC.Data[1908] := 37.042;
   Prof_FEC.Data[1909] := 34.325;
   Prof_FEC.Data[1910] := 37.025;
   Prof_FEC.Data[1911] := 37.715;
   Prof_FEC.Data[1912] := 36.962;
   Prof_FEC.Data[1913] := 38.014;
   Prof_FEC.Data[1914] := 39.643;
   Prof_FEC.Data[1915] := 39.128;
   Prof_FEC.Data[1916] := 38.145;
   Prof_FEC.Data[1917] := 36.441;
   Prof_FEC.Data[1918] := 38.582;
   Prof_FEC.Data[1919] := 38.282;
   Prof_FEC.Data[1920] := 40.068;
   Prof_FEC.Data[1921] := 39.526;
   Prof_FEC.Data[1922] := 37.093;
   Prof_FEC.Data[1923] := 38.541;
   Prof_FEC.Data[1924] := 39.449;
   Prof_FEC.Data[1925] := 36.215;
   Prof_FEC.Data[1926] := 40.342;
   Prof_FEC.Data[1927] := 38.674;
   Prof_FEC.Data[1928] := 43.669;
   Prof_FEC.Data[1929] := 43.344;
   Prof_FEC.Data[1930] := 39.974;
   Prof_FEC.Data[1931] := 39.155;
   Prof_FEC.Data[1932] := 40.612;
   Prof_FEC.Data[1933] := 40.175;
   Prof_FEC.Data[1934] := 38.762;
   Prof_FEC.Data[1935] := 38.989;
   Prof_FEC.Data[1936] := 37.221;
   Prof_FEC.Data[1937] := 39.139;
   Prof_FEC.Data[1938] := 37.041;
   Prof_FEC.Data[1939] := 36.046;
   Prof_FEC.Data[1940] := 193.82;
   Prof_FEC.Data[1941] := 192.2;
   Prof_FEC.Data[1942] := 217.86;
   Prof_FEC.Data[1943] := 247.64;
   Prof_FEC.Data[1944] := 294.95;
   Prof_FEC.Data[1945] := 391.4;
   Prof_FEC.Data[1946] := 387.89;
   Prof_FEC.Data[1947] := 368.66;
   Prof_FEC.Data[1948] := 430.8;
   Prof_FEC.Data[1949] := 490.93;
   Prof_FEC.Data[1950] := 482.08;
   Prof_FEC.Data[1951] := 460.0;
   Prof_FEC.Data[1952] := 474.05;
   Prof_FEC.Data[1953] := 446.66;
   Prof_FEC.Data[1954] := 472.69;
   Prof_FEC.Data[1955] := 494.72;
   Prof_FEC.Data[1956] := 512.99;
   Prof_FEC.Data[1957] := 569.57;
   Prof_FEC.Data[1958] := 580.45;
   Prof_FEC.Data[1959] := 536.62;
   Prof_FEC.Data[1960] := 558.75;
   Prof_FEC.Data[1961] := 634.5;
   Prof_FEC.Data[1962] := 601.98;
   Prof_FEC.Data[1963] := 555.79;
   Prof_FEC.Data[1964] := 624.92;
   Prof_FEC.Data[1965] := 592.41;
   Prof_FEC.Data[1966] := 593.05;
   Prof_FEC.Data[1967] := 551.63;
   Prof_FEC.Data[1968] := 565.73;
   Prof_FEC.Data[1969] := 558.75;
   Prof_FEC.Data[1970] := 449.33;
   Prof_FEC.Data[1971] := 515.97;
   Prof_FEC.Data[1972] := 526.67;
   Prof_FEC.Data[1973] := 554.83;
   Prof_FEC.Data[1974] := 540.44;
   Prof_FEC.Data[1975] := 530.72;
   Prof_FEC.Data[1976] := 578.96;
   Prof_FEC.Data[1977] := 484.25;
   Prof_FEC.Data[1978] := 501.75;
   Prof_FEC.Data[1979] := 559.58;
   Prof_FEC.Data[1980] := 609.51;
   Prof_FEC.Data[1981] := 526.54;
   Prof_FEC.Data[1982] := 628.28;
   Prof_FEC.Data[1983] := 601.04;
   Prof_FEC.Data[1984] := 703.39;
   Prof_FEC.Data[1985] := 736.82;
   Prof_FEC.Data[1986] := 705.86;
   Prof_FEC.Data[1987] := 598.33;
   Prof_FEC.Data[1988] := 406.93;
   Prof_FEC.Data[1989] := 376.83;
   Prof_FEC.Data[1990] := 335.94;
   Prof_FEC.Data[1991] := 290.98;
   Prof_FEC.Data[1992] := 259.16;
   Prof_FEC.Data[1993] := 233.18;
   Prof_FEC.Data[1994] := 234.94;
   Prof_FEC.Data[1995] := 228.15;
   Prof_FEC.Data[1996] := 39.185;
   Prof_FEC.Data[1997] := 42.393;
   Prof_FEC.Data[1998] := 39.447;
   Prof_FEC.Data[1999] := 41.223;
   Prof_FEC.Data[2000] := 39.335;
   Prof_FEC.Data[2001] := 39.733;
   Prof_FEC.Data[2002] := 39.726;
   Prof_FEC.Data[2003] := 37.35;
   Prof_FEC.Data[2004] := 41.837;
   Prof_FEC.Data[2005] := 40.503;
   Prof_FEC.Data[2006] := 42.564;
   Prof_FEC.Data[2007] := 42.32;
   Prof_FEC.Data[2008] := 39.68;
   Prof_FEC.Data[2009] := 40.437;
   Prof_FEC.Data[2010] := 38.661;
   Prof_FEC.Data[2011] := 42.524;
   Prof_FEC.Data[2012] := 44.017;
   Prof_FEC.Data[2013] := 46.97;
   Prof_FEC.Data[2014] := 42.377;
   Prof_FEC.Data[2015] := 41.117;
   Prof_FEC.Data[2016] := 40.641;
   Prof_FEC.Data[2017] := 39.567;
   Prof_FEC.Data[2018] := 39.482;
   Prof_FEC.Data[2019] := 41.446;
   Prof_FEC.Data[2020] := 42.224;
   Prof_FEC.Data[2021] := 39.902;
   Prof_FEC.Data[2022] := 41.824;
   Prof_FEC.Data[2023] := 40.105;
   Prof_FEC.Data[2024] := 39.152;
   Prof_FEC.Data[2025] := 39.833;
   Prof_FEC.Data[2026] := 38.9;
   Prof_FEC.Data[2027] := 38.155;
   Prof_FEC.Data[2028] := 39.073;
   Prof_FEC.Data[2029] := 37.463;
   Prof_FEC.Data[2030] := 38.622;
   Prof_FEC.Data[2031] := 40.674;
   Prof_FEC.Data[2032] := 37.4;
   Prof_FEC.Data[2033] := 39.629;
   Prof_FEC.Data[2034] := 38.555;
   Prof_FEC.Data[2035] := 38.399;
   Prof_FEC.Data[2036] := 224.42;
   Prof_FEC.Data[2037] := 235.5;
   Prof_FEC.Data[2038] := 249.26;
   Prof_FEC.Data[2039] := 260.75;
   Prof_FEC.Data[2040] := 308.76;
   Prof_FEC.Data[2041] := 342.15;
   Prof_FEC.Data[2042] := 405.73;
   Prof_FEC.Data[2043] := 409.2;
   Prof_FEC.Data[2044] := 516.04;
   Prof_FEC.Data[2045] := 511.48;
   Prof_FEC.Data[2046] := 557.53;
   Prof_FEC.Data[2047] := 560.93;
   Prof_FEC.Data[2048] := 602.03;
   Prof_FEC.Data[2049] := 592.48;
   Prof_FEC.Data[2050] := 646.3;
   Prof_FEC.Data[2051] := 642.75;
   Prof_FEC.Data[2052] := 675.39;
   Prof_FEC.Data[2053] := 623.97;
   Prof_FEC.Data[2054] := 662.34;
   Prof_FEC.Data[2055] := 618.73;
   Prof_FEC.Data[2056] := 612.82;
   Prof_FEC.Data[2057] := 650.97;
   Prof_FEC.Data[2058] := 654.21;
   Prof_FEC.Data[2059] := 623.09;
   Prof_FEC.Data[2060] := 685.24;
   Prof_FEC.Data[2061] := 668.59;
   Prof_FEC.Data[2062] := 592.28;
   Prof_FEC.Data[2063] := 624.0;
   Prof_FEC.Data[2064] := 580.57;
   Prof_FEC.Data[2065] := 574.97;
   Prof_FEC.Data[2066] := 527.38;
   Prof_FEC.Data[2067] := 567.32;
   Prof_FEC.Data[2068] := 624.53;
   Prof_FEC.Data[2069] := 624.09;
   Prof_FEC.Data[2070] := 562.75;
   Prof_FEC.Data[2071] := 564.57;
   Prof_FEC.Data[2072] := 679.67;
   Prof_FEC.Data[2073] := 583.91;
   Prof_FEC.Data[2074] := 625.04;
   Prof_FEC.Data[2075] := 629.27;
   Prof_FEC.Data[2076] := 514.4;
   Prof_FEC.Data[2077] := 532.19;
   Prof_FEC.Data[2078] := 511.96;
   Prof_FEC.Data[2079] := 638.49;
   Prof_FEC.Data[2080] := 705.27;
   Prof_FEC.Data[2081] := 676.97;
   Prof_FEC.Data[2082] := 651.79;
   Prof_FEC.Data[2083] := 569.17;
   Prof_FEC.Data[2084] := 394.69;
   Prof_FEC.Data[2085] := 299.41;
   Prof_FEC.Data[2086] := 326.34;
   Prof_FEC.Data[2087] := 219.52;
   Prof_FEC.Data[2088] := 235.54;
   Prof_FEC.Data[2089] := 220.04;
   Prof_FEC.Data[2090] := 228.57;
   Prof_FEC.Data[2091] := 235.56;
   Prof_FEC.Data[2092] := 40.149;
   Prof_FEC.Data[2093] := 40.868;
   Prof_FEC.Data[2094] := 39.459;
   Prof_FEC.Data[2095] := 39.515;
   Prof_FEC.Data[2096] := 39.442;
   Prof_FEC.Data[2097] := 37.65;
   Prof_FEC.Data[2098] := 37.295;
   Prof_FEC.Data[2099] := 40.733;
   Prof_FEC.Data[2100] := 40.8;
   Prof_FEC.Data[2101] := 41.663;
   Prof_FEC.Data[2102] := 37.61;
   Prof_FEC.Data[2103] := 39.926;
   Prof_FEC.Data[2104] := 39.163;
   Prof_FEC.Data[2105] := 35.955;
   Prof_FEC.Data[2106] := 35.934;
   Prof_FEC.Data[2107] := 39.126;
   Prof_FEC.Data[2108] := 40.194;
   Prof_FEC.Data[2109] := 41.544;
   Prof_FEC.Data[2110] := 41.234;
   Prof_FEC.Data[2111] := 41.737;
   Prof_FEC.Data[2112] := 38.766;
   Prof_FEC.Data[2113] := 38.723;
   Prof_FEC.Data[2114] := 40.51;
   Prof_FEC.Data[2115] := 37.641;
   Prof_FEC.Data[2116] := 41.525;
   Prof_FEC.Data[2117] := 41.137;
   Prof_FEC.Data[2118] := 40.927;
   Prof_FEC.Data[2119] := 40.192;
   Prof_FEC.Data[2120] := 37.106;
   Prof_FEC.Data[2121] := 39.85;
   Prof_FEC.Data[2122] := 36.575;
   Prof_FEC.Data[2123] := 37.058;
   Prof_FEC.Data[2124] := 39.896;
   Prof_FEC.Data[2125] := 40.897;
   Prof_FEC.Data[2126] := 43.914;
   Prof_FEC.Data[2127] := 40.6;
   Prof_FEC.Data[2128] := 41.582;
   Prof_FEC.Data[2129] := 39.669;
   Prof_FEC.Data[2130] := 38.379;
   Prof_FEC.Data[2131] := 41.238;
   Prof_FEC.Data[2132] := 235.13;
   Prof_FEC.Data[2133] := 254.25;
   Prof_FEC.Data[2134] := 277.01;
   Prof_FEC.Data[2135] := 295.65;
   Prof_FEC.Data[2136] := 313.85;
   Prof_FEC.Data[2137] := 319.42;
   Prof_FEC.Data[2138] := 394.86;
   Prof_FEC.Data[2139] := 420.7;
   Prof_FEC.Data[2140] := 509.42;
   Prof_FEC.Data[2141] := 568.61;
   Prof_FEC.Data[2142] := 561.85;
   Prof_FEC.Data[2143] := 583.5;
   Prof_FEC.Data[2144] := 558.3;
   Prof_FEC.Data[2145] := 575.52;
   Prof_FEC.Data[2146] := 572.25;
   Prof_FEC.Data[2147] := 624.27;
   Prof_FEC.Data[2148] := 582.19;
   Prof_FEC.Data[2149] := 576.46;
   Prof_FEC.Data[2150] := 581.85;
   Prof_FEC.Data[2151] := 630.38;
   Prof_FEC.Data[2152] := 620.29;
   Prof_FEC.Data[2153] := 694.82;
   Prof_FEC.Data[2154] := 608.55;
   Prof_FEC.Data[2155] := 686.71;
   Prof_FEC.Data[2156] := 623.0;
   Prof_FEC.Data[2157] := 632.32;
   Prof_FEC.Data[2158] := 673.48;
   Prof_FEC.Data[2159] := 711.17;
   Prof_FEC.Data[2160] := 627.62;
   Prof_FEC.Data[2161] := 569.63;
   Prof_FEC.Data[2162] := 548.46;
   Prof_FEC.Data[2163] := 587.86;
   Prof_FEC.Data[2164] := 647.51;
   Prof_FEC.Data[2165] := 685.8;
   Prof_FEC.Data[2166] := 599.33;
   Prof_FEC.Data[2167] := 604.13;
   Prof_FEC.Data[2168] := 676.56;
   Prof_FEC.Data[2169] := 710.74;
   Prof_FEC.Data[2170] := 731.32;
   Prof_FEC.Data[2171] := 586.77;
   Prof_FEC.Data[2172] := 702.4;
   Prof_FEC.Data[2173] := 671.91;
   Prof_FEC.Data[2174] := 641.13;
   Prof_FEC.Data[2175] := 684.0;
   Prof_FEC.Data[2176] := 747.29;
   Prof_FEC.Data[2177] := 656.66;
   Prof_FEC.Data[2178] := 625.43;
   Prof_FEC.Data[2179] := 548.57;
   Prof_FEC.Data[2180] := 377.64;
   Prof_FEC.Data[2181] := 354.03;
   Prof_FEC.Data[2182] := 306.94;
   Prof_FEC.Data[2183] := 259.26;
   Prof_FEC.Data[2184] := 244.89;
   Prof_FEC.Data[2185] := 222.56;
   Prof_FEC.Data[2186] := 213.88;
   Prof_FEC.Data[2187] := 230.08;
   Prof_FEC.Data[2188] := 37.625;
   Prof_FEC.Data[2189] := 39.706;
   Prof_FEC.Data[2190] := 39.856;
   Prof_FEC.Data[2191] := 38.76;
   Prof_FEC.Data[2192] := 37.967;
   Prof_FEC.Data[2193] := 41.338;
   Prof_FEC.Data[2194] := 36.245;
   Prof_FEC.Data[2195] := 36.908;
   Prof_FEC.Data[2196] := 41.385;
   Prof_FEC.Data[2197] := 38.353;
   Prof_FEC.Data[2198] := 39.985;
   Prof_FEC.Data[2199] := 40.085;
   Prof_FEC.Data[2200] := 39.853;
   Prof_FEC.Data[2201] := 39.702;
   Prof_FEC.Data[2202] := 39.271;
   Prof_FEC.Data[2203] := 41.501;
   Prof_FEC.Data[2204] := 40.916;
   Prof_FEC.Data[2205] := 43.521;
   Prof_FEC.Data[2206] := 45.271;
   Prof_FEC.Data[2207] := 41.941;
   Prof_FEC.Data[2208] := 42.846;
   Prof_FEC.Data[2209] := 41.246;
   Prof_FEC.Data[2210] := 43.398;
   Prof_FEC.Data[2211] := 44.913;
   Prof_FEC.Data[2212] := 48.037;
   Prof_FEC.Data[2213] := 45.861;
   Prof_FEC.Data[2214] := 45.925;
   Prof_FEC.Data[2215] := 45.072;
   Prof_FEC.Data[2216] := 41.414;
   Prof_FEC.Data[2217] := 43.558;
   Prof_FEC.Data[2218] := 41.551;
   Prof_FEC.Data[2219] := 44.728;
   Prof_FEC.Data[2220] := 45.526;
   Prof_FEC.Data[2221] := 43.658;
   Prof_FEC.Data[2222] := 49.731;
   Prof_FEC.Data[2223] := 41.031;
   Prof_FEC.Data[2224] := 43.138;
   Prof_FEC.Data[2225] := 42.883;
   Prof_FEC.Data[2226] := 40.269;
   Prof_FEC.Data[2227] := 43.198;
   Prof_FEC.Data[2228] := 257.69;
   Prof_FEC.Data[2229] := 252.64;
   Prof_FEC.Data[2230] := 293.71;
   Prof_FEC.Data[2231] := 289.43;
   Prof_FEC.Data[2232] := 309.12;
   Prof_FEC.Data[2233] := 346.59;
   Prof_FEC.Data[2234] := 408.09;
   Prof_FEC.Data[2235] := 416.4;
   Prof_FEC.Data[2236] := 427.44;
   Prof_FEC.Data[2237] := 482.06;
   Prof_FEC.Data[2238] := 493.67;
   Prof_FEC.Data[2239] := 513.26;
   Prof_FEC.Data[2240] := 563.37;
   Prof_FEC.Data[2241] := 544.53;
   Prof_FEC.Data[2242] := 533.53;
   Prof_FEC.Data[2243] := 579.69;
   Prof_FEC.Data[2244] := 604.42;
   Prof_FEC.Data[2245] := 634.91;
   Prof_FEC.Data[2246] := 651.05;
   Prof_FEC.Data[2247] := 729.46;
   Prof_FEC.Data[2248] := 645.51;
   Prof_FEC.Data[2249] := 638.91;
   Prof_FEC.Data[2250] := 702.06;
   Prof_FEC.Data[2251] := 618.28;
   Prof_FEC.Data[2252] := 674.66;
   Prof_FEC.Data[2253] := 710.39;
   Prof_FEC.Data[2254] := 621.97;
   Prof_FEC.Data[2255] := 669.38;
   Prof_FEC.Data[2256] := 577.34;
   Prof_FEC.Data[2257] := 532.8;
   Prof_FEC.Data[2258] := 537.44;
   Prof_FEC.Data[2259] := 542.37;
   Prof_FEC.Data[2260] := 571.76;
   Prof_FEC.Data[2261] := 683.16;
   Prof_FEC.Data[2262] := 685.78;
   Prof_FEC.Data[2263] := 631.45;
   Prof_FEC.Data[2264] := 614.98;
   Prof_FEC.Data[2265] := 694.58;
   Prof_FEC.Data[2266] := 743.02;
   Prof_FEC.Data[2267] := 652.92;
   Prof_FEC.Data[2268] := 609.2;
   Prof_FEC.Data[2269] := 601.05;
   Prof_FEC.Data[2270] := 658.85;
   Prof_FEC.Data[2271] := 667.55;
   Prof_FEC.Data[2272] := 648.92;
   Prof_FEC.Data[2273] := 670.93;
   Prof_FEC.Data[2274] := 649.32;
   Prof_FEC.Data[2275] := 572.5;
   Prof_FEC.Data[2276] := 438.03;
   Prof_FEC.Data[2277] := 321.35;
   Prof_FEC.Data[2278] := 297.72;
   Prof_FEC.Data[2279] := 241.73;
   Prof_FEC.Data[2280] := 190.53;
   Prof_FEC.Data[2281] := 239.59;
   Prof_FEC.Data[2282] := 200.77;
   Prof_FEC.Data[2283] := 206.95;
   Prof_FEC.Data[2284] := 36.327;
   Prof_FEC.Data[2285] := 37.27;
   Prof_FEC.Data[2286] := 40.076;
   Prof_FEC.Data[2287] := 36.925;
   Prof_FEC.Data[2288] := 38.447;
   Prof_FEC.Data[2289] := 38.796;
   Prof_FEC.Data[2290] := 38.338;
   Prof_FEC.Data[2291] := 38.877;
   Prof_FEC.Data[2292] := 42.055;
   Prof_FEC.Data[2293] := 41.328;
   Prof_FEC.Data[2294] := 37.811;
   Prof_FEC.Data[2295] := 40.273;
   Prof_FEC.Data[2296] := 41.941;
   Prof_FEC.Data[2297] := 36.625;
   Prof_FEC.Data[2298] := 40.387;
   Prof_FEC.Data[2299] := 37.695;
   Prof_FEC.Data[2300] := 37.043;
   Prof_FEC.Data[2301] := 37.809;
   Prof_FEC.Data[2302] := 39.725;
   Prof_FEC.Data[2303] := 39.566;
   Prof_FEC.Data[2304] := 34.174;
   Prof_FEC.Data[2305] := 37.001;
   Prof_FEC.Data[2306] := 33.239;
   Prof_FEC.Data[2307] := 36.974;
   Prof_FEC.Data[2308] := 36.857;
   Prof_FEC.Data[2309] := 39.56;
   Prof_FEC.Data[2310] := 37.75;
   Prof_FEC.Data[2311] := 39.281;
   Prof_FEC.Data[2312] := 36.839;
   Prof_FEC.Data[2313] := 37.152;
   Prof_FEC.Data[2314] := 34.875;
   Prof_FEC.Data[2315] := 37.79;
   Prof_FEC.Data[2316] := 38.958;
   Prof_FEC.Data[2317] := 41.528;
   Prof_FEC.Data[2318] := 40.256;
   Prof_FEC.Data[2319] := 41.093;
   Prof_FEC.Data[2320] := 39.965;
   Prof_FEC.Data[2321] := 38.859;
   Prof_FEC.Data[2322] := 38.828;
   Prof_FEC.Data[2323] := 35.894;
   Prof_FEC.Data[2324] := 224.45;
   Prof_FEC.Data[2325] := 217.46;
   Prof_FEC.Data[2326] := 237.71;
   Prof_FEC.Data[2327] := 235.91;
   Prof_FEC.Data[2328] := 203.75;
   Prof_FEC.Data[2329] := 171.87;
   Prof_FEC.Data[2330] := 193.96;
   Prof_FEC.Data[2331] := 211.98;
   Prof_FEC.Data[2332] := 265.56;
   Prof_FEC.Data[2333] := 293.61;
   Prof_FEC.Data[2334] := 356.48;
   Prof_FEC.Data[2335] := 296.16;
   Prof_FEC.Data[2336] := 239.99;
   Prof_FEC.Data[2337] := 240.98;
   Prof_FEC.Data[2338] := 226.85;
   Prof_FEC.Data[2339] := 241.87;
   Prof_FEC.Data[2340] := 296.2;
   Prof_FEC.Data[2341] := 301.72;
   Prof_FEC.Data[2342] := 312.27;
   Prof_FEC.Data[2343] := 312.42;
   Prof_FEC.Data[2344] := 309.22;
   Prof_FEC.Data[2345] := 288.76;
   Prof_FEC.Data[2346] := 278.53;
   Prof_FEC.Data[2347] := 327.11;
   Prof_FEC.Data[2348] := 333.6;
   Prof_FEC.Data[2349] := 331.02;
   Prof_FEC.Data[2350] := 328.16;
   Prof_FEC.Data[2351] := 289.76;
   Prof_FEC.Data[2352] := 230.07;
   Prof_FEC.Data[2353] := 255.29;
   Prof_FEC.Data[2354] := 223.53;
   Prof_FEC.Data[2355] := 251.04;
   Prof_FEC.Data[2356] := 279.0;
   Prof_FEC.Data[2357] := 268.64;
   Prof_FEC.Data[2358] := 257.97;
   Prof_FEC.Data[2359] := 259.77;
   Prof_FEC.Data[2360] := 258.49;
   Prof_FEC.Data[2361] := 261.25;
   Prof_FEC.Data[2362] := 262.9;
   Prof_FEC.Data[2363] := 294.85;
   Prof_FEC.Data[2364] := 338.78;
   Prof_FEC.Data[2365] := 310.97;
   Prof_FEC.Data[2366] := 277.43;
   Prof_FEC.Data[2367] := 245.88;
   Prof_FEC.Data[2368] := 172.5;
   Prof_FEC.Data[2369] := 147.98;
   Prof_FEC.Data[2370] := 156.82;
   Prof_FEC.Data[2371] := 169.61;
   Prof_FEC.Data[2372] := 188.81;
   Prof_FEC.Data[2373] := 214.44;
   Prof_FEC.Data[2374] := 239.7;
   Prof_FEC.Data[2375] := 232.19;
   Prof_FEC.Data[2376] := 239.56;
   Prof_FEC.Data[2377] := 265.15;
   Prof_FEC.Data[2378] := 266.85;
   Prof_FEC.Data[2379] := 261.83;
   Prof_FEC.Data[2380] := 40.12;
   Prof_FEC.Data[2381] := 39.756;
   Prof_FEC.Data[2382] := 38.605;
   Prof_FEC.Data[2383] := 39.715;
   Prof_FEC.Data[2384] := 40.061;
   Prof_FEC.Data[2385] := 42.635;
   Prof_FEC.Data[2386] := 42.345;
   Prof_FEC.Data[2387] := 42.462;
   Prof_FEC.Data[2388] := 38.428;
   Prof_FEC.Data[2389] := 39.944;
   Prof_FEC.Data[2390] := 39.827;
   Prof_FEC.Data[2391] := 40.869;
   Prof_FEC.Data[2392] := 42.761;
   Prof_FEC.Data[2393] := 41.705;
   Prof_FEC.Data[2394] := 42.226;
   Prof_FEC.Data[2395] := 41.609;
   Prof_FEC.Data[2396] := 38.408;
   Prof_FEC.Data[2397] := 42.936;
   Prof_FEC.Data[2398] := 41.558;
   Prof_FEC.Data[2399] := 43.679;
   Prof_FEC.Data[2400] := 42.934;
   Prof_FEC.Data[2401] := 42.545;
   Prof_FEC.Data[2402] := 43.235;
   Prof_FEC.Data[2403] := 43.985;
   Prof_FEC.Data[2404] := 42.215;
   Prof_FEC.Data[2405] := 41.381;
   Prof_FEC.Data[2406] := 40.238;
   Prof_FEC.Data[2407] := 41.23;
   Prof_FEC.Data[2408] := 40.436;
   Prof_FEC.Data[2409] := 42.721;
   Prof_FEC.Data[2410] := 39.709;
   Prof_FEC.Data[2411] := 37.926;
   Prof_FEC.Data[2412] := 37.583;
   Prof_FEC.Data[2413] := 40.382;
   Prof_FEC.Data[2414] := 39.725;
   Prof_FEC.Data[2415] := 38.076;
   Prof_FEC.Data[2416] := 42.448;
   Prof_FEC.Data[2417] := 42.433;
   Prof_FEC.Data[2418] := 42.415;
   Prof_FEC.Data[2419] := 43.262;
   Prof_FEC.Data[2420] := 252.9;
   Prof_FEC.Data[2421] := 258.77;
   Prof_FEC.Data[2422] := 230.08;
   Prof_FEC.Data[2423] := 278.82;
   Prof_FEC.Data[2424] := 283.5;
   Prof_FEC.Data[2425] := 285.06;
   Prof_FEC.Data[2426] := 310.87;
   Prof_FEC.Data[2427] := 291.38;
   Prof_FEC.Data[2428] := 258.89;
   Prof_FEC.Data[2429] := 260.71;
   Prof_FEC.Data[2430] := 253.9;
   Prof_FEC.Data[2431] := 205.53;
   Prof_FEC.Data[2432] := 194.49;
   Prof_FEC.Data[2433] := 171.39;
   Prof_FEC.Data[2434] := 166.6;
   Prof_FEC.Data[2435] := 169.22;
   Prof_FEC.Data[2436] := 147.75;
   Prof_FEC.Data[2437] := 172.26;
   Prof_FEC.Data[2438] := 160.41;
   Prof_FEC.Data[2439] := 182.01;
   Prof_FEC.Data[2440] := 185.16;
   Prof_FEC.Data[2441] := 180.01;
   Prof_FEC.Data[2442] := 179.76;
   Prof_FEC.Data[2443] := 177.94;
   Prof_FEC.Data[2444] := 141.81;
   Prof_FEC.Data[2445] := 144.72;
   Prof_FEC.Data[2446] := 148.99;
   Prof_FEC.Data[2447] := 145.68;
   Prof_FEC.Data[2448] := 173.25;
   Prof_FEC.Data[2449] := 170.52;
   Prof_FEC.Data[2450] := 194.46;
   Prof_FEC.Data[2451] := 177.35;
   Prof_FEC.Data[2452] := 160.94;
   Prof_FEC.Data[2453] := 133.09;
   Prof_FEC.Data[2454] := 150.92;
   Prof_FEC.Data[2455] := 144.04;
   Prof_FEC.Data[2456] := 142.01;
   Prof_FEC.Data[2457] := 161.03;
   Prof_FEC.Data[2458] := 148.5;
   Prof_FEC.Data[2459] := 155.39;
   Prof_FEC.Data[2460] := 140.27;
   Prof_FEC.Data[2461] := 113.58;
   Prof_FEC.Data[2462] := 121.99;
   Prof_FEC.Data[2463] := 132.11;
   Prof_FEC.Data[2464] := 146.15;
   Prof_FEC.Data[2465] := 195.49;
   Prof_FEC.Data[2466] := 201.02;
   Prof_FEC.Data[2467] := 234.68;
   Prof_FEC.Data[2468] := 240.62;
   Prof_FEC.Data[2469] := 243.9;
   Prof_FEC.Data[2470] := 274.05;
   Prof_FEC.Data[2471] := 289.96;
   Prof_FEC.Data[2472] := 270.63;
   Prof_FEC.Data[2473] := 304.79;
   Prof_FEC.Data[2474] := 259.0;
   Prof_FEC.Data[2475] := 318.96;
   Prof_FEC.Data[2476] := 44.115;
   Prof_FEC.Data[2477] := 39.738;
   Prof_FEC.Data[2478] := 43.809;
   Prof_FEC.Data[2479] := 41.988;
   Prof_FEC.Data[2480] := 46.866;
   Prof_FEC.Data[2481] := 48.766;
   Prof_FEC.Data[2482] := 45.771;
   Prof_FEC.Data[2483] := 48.748;
   Prof_FEC.Data[2484] := 44.961;
   Prof_FEC.Data[2485] := 42.633;
   Prof_FEC.Data[2486] := 43.713;
   Prof_FEC.Data[2487] := 43.275;
   Prof_FEC.Data[2488] := 45.749;
   Prof_FEC.Data[2489] := 46.329;
   Prof_FEC.Data[2490] := 47.598;
   Prof_FEC.Data[2491] := 47.749;
   Prof_FEC.Data[2492] := 42.217;
   Prof_FEC.Data[2493] := 41.669;
   Prof_FEC.Data[2494] := 41.843;
   Prof_FEC.Data[2495] := 41.553;
   Prof_FEC.Data[2496] := 50.0;
   Prof_FEC.Data[2497] := 47.49;
   Prof_FEC.Data[2498] := 49.039;
   Prof_FEC.Data[2499] := 50.0;
   Prof_FEC.Data[2500] := 45.754;
   Prof_FEC.Data[2501] := 46.008;
   Prof_FEC.Data[2502] := 43.465;
   Prof_FEC.Data[2503] := 49.027;
   Prof_FEC.Data[2504] := 49.802;
   Prof_FEC.Data[2505] := 49.151;
   Prof_FEC.Data[2506] := 48.215;
   Prof_FEC.Data[2507] := 50.0;
   Prof_FEC.Data[2508] := 45.661;
   Prof_FEC.Data[2509] := 44.445;
   Prof_FEC.Data[2510] := 47.22;
   Prof_FEC.Data[2511] := 48.092;
   Prof_FEC.Data[2512] := 50.0;
   Prof_FEC.Data[2513] := 50.0;
   Prof_FEC.Data[2514] := 50.0;
   Prof_FEC.Data[2515] := 50.0;
   Prof_FEC.Data[2516] := 339.2;
   Prof_FEC.Data[2517] := 364.48;
   Prof_FEC.Data[2518] := 324.98;
   Prof_FEC.Data[2519] := 374.0;
   Prof_FEC.Data[2520] := 386.08;
   Prof_FEC.Data[2521] := 403.73;
   Prof_FEC.Data[2522] := 426.53;
   Prof_FEC.Data[2523] := 512.36;
   Prof_FEC.Data[2524] := 567.1;
   Prof_FEC.Data[2525] := 531.37;
   Prof_FEC.Data[2526] := 601.66;
   Prof_FEC.Data[2527] := 652.0;
   Prof_FEC.Data[2528] := 627.37;
   Prof_FEC.Data[2529] := 609.12;
   Prof_FEC.Data[2530] := 585.73;
   Prof_FEC.Data[2531] := 668.51;
   Prof_FEC.Data[2532] := 704.71;
   Prof_FEC.Data[2533] := 721.29;
   Prof_FEC.Data[2534] := 712.02;
   Prof_FEC.Data[2535] := 687.72;
   Prof_FEC.Data[2536] := 700.13;
   Prof_FEC.Data[2537] := 672.9;
   Prof_FEC.Data[2538] := 625.86;
   Prof_FEC.Data[2539] := 670.48;
   Prof_FEC.Data[2540] := 703.7;
   Prof_FEC.Data[2541] := 669.85;
   Prof_FEC.Data[2542] := 615.24;
   Prof_FEC.Data[2543] := 629.93;
   Prof_FEC.Data[2544] := 588.8;
   Prof_FEC.Data[2545] := 598.6;
   Prof_FEC.Data[2546] := 686.68;
   Prof_FEC.Data[2547] := 635.77;
   Prof_FEC.Data[2548] := 633.96;
   Prof_FEC.Data[2549] := 703.11;
   Prof_FEC.Data[2550] := 769.4;
   Prof_FEC.Data[2551] := 750.12;
   Prof_FEC.Data[2552] := 739.25;
   Prof_FEC.Data[2553] := 728.14;
   Prof_FEC.Data[2554] := 680.53;
   Prof_FEC.Data[2555] := 640.2;
   Prof_FEC.Data[2556] := 681.49;
   Prof_FEC.Data[2557] := 598.34;
   Prof_FEC.Data[2558] := 624.34;
   Prof_FEC.Data[2559] := 623.13;
   Prof_FEC.Data[2560] := 613.34;
   Prof_FEC.Data[2561] := 752.41;
   Prof_FEC.Data[2562] := 709.74;
   Prof_FEC.Data[2563] := 533.3;
   Prof_FEC.Data[2564] := 535.69;
   Prof_FEC.Data[2565] := 435.98;
   Prof_FEC.Data[2566] := 386.46;
   Prof_FEC.Data[2567] := 329.99;
   Prof_FEC.Data[2568] := 258.46;
   Prof_FEC.Data[2569] := 255.41;
   Prof_FEC.Data[2570] := 234.29;
   Prof_FEC.Data[2571] := 234.45;
   Prof_FEC.Data[2572] := 46.995;
   Prof_FEC.Data[2573] := 47.695;
   Prof_FEC.Data[2574] := 50.0;
   Prof_FEC.Data[2575] := 45.388;
   Prof_FEC.Data[2576] := 41.361;
   Prof_FEC.Data[2577] := 42.875;
   Prof_FEC.Data[2578] := 41.115;
   Prof_FEC.Data[2579] := 41.019;
   Prof_FEC.Data[2580] := 44.481;
   Prof_FEC.Data[2581] := 44.473;
   Prof_FEC.Data[2582] := 43.889;
   Prof_FEC.Data[2583] := 41.192;
   Prof_FEC.Data[2584] := 42.128;
   Prof_FEC.Data[2585] := 39.721;
   Prof_FEC.Data[2586] := 41.337;
   Prof_FEC.Data[2587] := 42.621;
   Prof_FEC.Data[2588] := 47.047;
   Prof_FEC.Data[2589] := 45.643;
   Prof_FEC.Data[2590] := 45.107;
   Prof_FEC.Data[2591] := 43.691;
   Prof_FEC.Data[2592] := 42.815;
   Prof_FEC.Data[2593] := 42.874;
   Prof_FEC.Data[2594] := 42.01;
   Prof_FEC.Data[2595] := 45.133;
   Prof_FEC.Data[2596] := 50.0;
   Prof_FEC.Data[2597] := 50.0;
   Prof_FEC.Data[2598] := 47.517;
   Prof_FEC.Data[2599] := 47.801;
   Prof_FEC.Data[2600] := 43.685;
   Prof_FEC.Data[2601] := 46.313;
   Prof_FEC.Data[2602] := 43.935;
   Prof_FEC.Data[2603] := 42.233;
   Prof_FEC.Data[2604] := 44.825;
   Prof_FEC.Data[2605] := 43.911;
   Prof_FEC.Data[2606] := 47.375;
   Prof_FEC.Data[2607] := 47.055;
   Prof_FEC.Data[2608] := 39.196;
   Prof_FEC.Data[2609] := 42.232;
   Prof_FEC.Data[2610] := 40.752;
   Prof_FEC.Data[2611] := 44.079;
   Prof_FEC.Data[2612] := 272.82;
   Prof_FEC.Data[2613] := 311.87;
   Prof_FEC.Data[2614] := 321.98;
   Prof_FEC.Data[2615] := 351.42;
   Prof_FEC.Data[2616] := 358.37;
   Prof_FEC.Data[2617] := 401.28;
   Prof_FEC.Data[2618] := 412.29;
   Prof_FEC.Data[2619] := 462.34;
   Prof_FEC.Data[2620] := 458.83;
   Prof_FEC.Data[2621] := 512.11;
   Prof_FEC.Data[2622] := 514.15;
   Prof_FEC.Data[2623] := 533.25;
   Prof_FEC.Data[2624] := 510.11;
   Prof_FEC.Data[2625] := 559.1;
   Prof_FEC.Data[2626] := 542.46;
   Prof_FEC.Data[2627] := 537.49;
   Prof_FEC.Data[2628] := 610.84;
   Prof_FEC.Data[2629] := 702.04;
   Prof_FEC.Data[2630] := 592.96;
   Prof_FEC.Data[2631] := 583.1;
   Prof_FEC.Data[2632] := 605.37;
   Prof_FEC.Data[2633] := 602.11;
   Prof_FEC.Data[2634] := 606.12;
   Prof_FEC.Data[2635] := 589.45;
   Prof_FEC.Data[2636] := 641.26;
   Prof_FEC.Data[2637] := 579.18;
   Prof_FEC.Data[2638] := 667.93;
   Prof_FEC.Data[2639] := 574.69;
   Prof_FEC.Data[2640] := 552.23;
   Prof_FEC.Data[2641] := 588.88;
   Prof_FEC.Data[2642] := 540.01;
   Prof_FEC.Data[2643] := 657.66;
   Prof_FEC.Data[2644] := 555.28;
   Prof_FEC.Data[2645] := 625.65;
   Prof_FEC.Data[2646] := 648.6;
   Prof_FEC.Data[2647] := 583.84;
   Prof_FEC.Data[2648] := 596.51;
   Prof_FEC.Data[2649] := 627.0;
   Prof_FEC.Data[2650] := 665.64;
   Prof_FEC.Data[2651] := 608.97;
   Prof_FEC.Data[2652] := 599.05;
   Prof_FEC.Data[2653] := 587.17;
   Prof_FEC.Data[2654] := 575.06;
   Prof_FEC.Data[2655] := 563.93;
   Prof_FEC.Data[2656] := 667.8;
   Prof_FEC.Data[2657] := 696.57;
   Prof_FEC.Data[2658] := 635.1;
   Prof_FEC.Data[2659] := 529.2;
   Prof_FEC.Data[2660] := 375.39;
   Prof_FEC.Data[2661] := 383.19;
   Prof_FEC.Data[2662] := 307.15;
   Prof_FEC.Data[2663] := 284.07;
   Prof_FEC.Data[2664] := 232.46;
   Prof_FEC.Data[2665] := 238.11;
   Prof_FEC.Data[2666] := 241.84;
   Prof_FEC.Data[2667] := 241.53;
   Prof_FEC.Data[2668] := 42.167;
   Prof_FEC.Data[2669] := 43.655;
   Prof_FEC.Data[2670] := 45.533;
   Prof_FEC.Data[2671] := 44.144;
   Prof_FEC.Data[2672] := 45.333;
   Prof_FEC.Data[2673] := 42.745;
   Prof_FEC.Data[2674] := 42.286;
   Prof_FEC.Data[2675] := 43.766;
   Prof_FEC.Data[2676] := 46.933;
   Prof_FEC.Data[2677] := 49.234;
   Prof_FEC.Data[2678] := 48.251;
   Prof_FEC.Data[2679] := 46.37;
   Prof_FEC.Data[2680] := 46.899;
   Prof_FEC.Data[2681] := 44.353;
   Prof_FEC.Data[2682] := 42.737;
   Prof_FEC.Data[2683] := 43.839;
   Prof_FEC.Data[2684] := 46.96;
   Prof_FEC.Data[2685] := 48.365;
   Prof_FEC.Data[2686] := 45.428;
   Prof_FEC.Data[2687] := 41.526;
   Prof_FEC.Data[2688] := 40.75;
   Prof_FEC.Data[2689] := 39.736;
   Prof_FEC.Data[2690] := 39.381;
   Prof_FEC.Data[2691] := 43.269;
   Prof_FEC.Data[2692] := 47.978;
   Prof_FEC.Data[2693] := 47.416;
   Prof_FEC.Data[2694] := 46.652;
   Prof_FEC.Data[2695] := 46.741;
   Prof_FEC.Data[2696] := 46.392;
   Prof_FEC.Data[2697] := 47.044;
   Prof_FEC.Data[2698] := 46.094;
   Prof_FEC.Data[2699] := 48.199;
   Prof_FEC.Data[2700] := 49.216;
   Prof_FEC.Data[2701] := 50.0;
   Prof_FEC.Data[2702] := 50.0;
   Prof_FEC.Data[2703] := 49.961;
   Prof_FEC.Data[2704] := 46.793;
   Prof_FEC.Data[2705] := 49.426;
   Prof_FEC.Data[2706] := 48.916;
   Prof_FEC.Data[2707] := 44.756;
   Prof_FEC.Data[2708] := 342.89;
   Prof_FEC.Data[2709] := 363.26;
   Prof_FEC.Data[2710] := 324.39;
   Prof_FEC.Data[2711] := 381.35;
   Prof_FEC.Data[2712] := 392.15;
   Prof_FEC.Data[2713] := 385.61;
   Prof_FEC.Data[2714] := 478.19;
   Prof_FEC.Data[2715] := 438.93;
   Prof_FEC.Data[2716] := 490.47;
   Prof_FEC.Data[2717] := 497.26;
   Prof_FEC.Data[2718] := 518.51;
   Prof_FEC.Data[2719] := 547.37;
   Prof_FEC.Data[2720] := 567.33;
   Prof_FEC.Data[2721] := 670.74;
   Prof_FEC.Data[2722] := 681.12;
   Prof_FEC.Data[2723] := 705.2;
   Prof_FEC.Data[2724] := 745.75;
   Prof_FEC.Data[2725] := 736.62;
   Prof_FEC.Data[2726] := 756.66;
   Prof_FEC.Data[2727] := 734.33;
   Prof_FEC.Data[2728] := 702.68;
   Prof_FEC.Data[2729] := 655.5;
   Prof_FEC.Data[2730] := 633.0;
   Prof_FEC.Data[2731] := 669.24;
   Prof_FEC.Data[2732] := 696.36;
   Prof_FEC.Data[2733] := 756.14;
   Prof_FEC.Data[2734] := 752.19;
   Prof_FEC.Data[2735] := 715.55;
   Prof_FEC.Data[2736] := 673.37;
   Prof_FEC.Data[2737] := 627.47;
   Prof_FEC.Data[2738] := 667.26;
   Prof_FEC.Data[2739] := 600.82;
   Prof_FEC.Data[2740] := 654.9;
   Prof_FEC.Data[2741] := 693.14;
   Prof_FEC.Data[2742] := 666.96;
   Prof_FEC.Data[2743] := 689.09;
   Prof_FEC.Data[2744] := 819.31;
   Prof_FEC.Data[2745] := 730.7;
   Prof_FEC.Data[2746] := 690.43;
   Prof_FEC.Data[2747] := 746.8;
   Prof_FEC.Data[2748] := 741.29;
   Prof_FEC.Data[2749] := 784.64;
   Prof_FEC.Data[2750] := 771.77;
   Prof_FEC.Data[2751] := 777.16;
   Prof_FEC.Data[2752] := 794.13;
   Prof_FEC.Data[2753] := 793.14;
   Prof_FEC.Data[2754] := 756.83;
   Prof_FEC.Data[2755] := 637.21;
   Prof_FEC.Data[2756] := 524.4;
   Prof_FEC.Data[2757] := 450.05;
   Prof_FEC.Data[2758] := 364.57;
   Prof_FEC.Data[2759] := 347.15;
   Prof_FEC.Data[2760] := 317.26;
   Prof_FEC.Data[2761] := 303.49;
   Prof_FEC.Data[2762] := 264.08;
   Prof_FEC.Data[2763] := 274.49;
   Prof_FEC.Data[2764] := 46.506;
   Prof_FEC.Data[2765] := 49.09;
   Prof_FEC.Data[2766] := 47.574;
   Prof_FEC.Data[2767] := 45.439;
   Prof_FEC.Data[2768] := 43.325;
   Prof_FEC.Data[2769] := 43.344;
   Prof_FEC.Data[2770] := 40.917;
   Prof_FEC.Data[2771] := 40.831;
   Prof_FEC.Data[2772] := 44.063;
   Prof_FEC.Data[2773] := 46.866;
   Prof_FEC.Data[2774] := 45.695;
   Prof_FEC.Data[2775] := 49.472;
   Prof_FEC.Data[2776] := 41.684;
   Prof_FEC.Data[2777] := 41.715;
   Prof_FEC.Data[2778] := 40.578;
   Prof_FEC.Data[2779] := 42.069;
   Prof_FEC.Data[2780] := 43.923;
   Prof_FEC.Data[2781] := 43.474;
   Prof_FEC.Data[2782] := 42.6;
   Prof_FEC.Data[2783] := 43.803;
   Prof_FEC.Data[2784] := 40.696;
   Prof_FEC.Data[2785] := 42.002;
   Prof_FEC.Data[2786] := 43.003;
   Prof_FEC.Data[2787] := 42.449;
   Prof_FEC.Data[2788] := 47.401;
   Prof_FEC.Data[2789] := 46.432;
   Prof_FEC.Data[2790] := 44.867;
   Prof_FEC.Data[2791] := 42.886;
   Prof_FEC.Data[2792] := 40.15;
   Prof_FEC.Data[2793] := 39.287;
   Prof_FEC.Data[2794] := 39.071;
   Prof_FEC.Data[2795] := 41.296;
   Prof_FEC.Data[2796] := 41.254;
   Prof_FEC.Data[2797] := 42.83;
   Prof_FEC.Data[2798] := 43.972;
   Prof_FEC.Data[2799] := 45.19;
   Prof_FEC.Data[2800] := 42.83;
   Prof_FEC.Data[2801] := 41.537;
   Prof_FEC.Data[2802] := 42.678;
   Prof_FEC.Data[2803] := 40.895;
   Prof_FEC.Data[2804] := 269.25;
   Prof_FEC.Data[2805] := 262.03;
   Prof_FEC.Data[2806] := 287.58;
   Prof_FEC.Data[2807] := 301.03;
   Prof_FEC.Data[2808] := 317.1;
   Prof_FEC.Data[2809] := 334.03;
   Prof_FEC.Data[2810] := 372.77;
   Prof_FEC.Data[2811] := 437.99;
   Prof_FEC.Data[2812] := 498.82;
   Prof_FEC.Data[2813] := 539.88;
   Prof_FEC.Data[2814] := 508.56;
   Prof_FEC.Data[2815] := 507.63;
   Prof_FEC.Data[2816] := 546.6;
   Prof_FEC.Data[2817] := 513.02;
   Prof_FEC.Data[2818] := 569.37;
   Prof_FEC.Data[2819] := 550.71;
   Prof_FEC.Data[2820] := 517.09;
   Prof_FEC.Data[2821] := 667.2;
   Prof_FEC.Data[2822] := 610.46;
   Prof_FEC.Data[2823] := 638.99;
   Prof_FEC.Data[2824] := 639.16;
   Prof_FEC.Data[2825] := 640.79;
   Prof_FEC.Data[2826] := 651.56;
   Prof_FEC.Data[2827] := 628.84;
   Prof_FEC.Data[2828] := 689.05;
   Prof_FEC.Data[2829] := 739.97;
   Prof_FEC.Data[2830] := 664.63;
   Prof_FEC.Data[2831] := 691.3;
   Prof_FEC.Data[2832] := 632.1;
   Prof_FEC.Data[2833] := 628.62;
   Prof_FEC.Data[2834] := 657.73;
   Prof_FEC.Data[2835] := 637.31;
   Prof_FEC.Data[2836] := 700.92;
   Prof_FEC.Data[2837] := 693.45;
   Prof_FEC.Data[2838] := 629.24;
   Prof_FEC.Data[2839] := 701.89;
   Prof_FEC.Data[2840] := 700.03;
   Prof_FEC.Data[2841] := 656.25;
   Prof_FEC.Data[2842] := 631.63;
   Prof_FEC.Data[2843] := 623.56;
   Prof_FEC.Data[2844] := 564.38;
   Prof_FEC.Data[2845] := 623.48;
   Prof_FEC.Data[2846] := 610.23;
   Prof_FEC.Data[2847] := 552.48;
   Prof_FEC.Data[2848] := 572.59;
   Prof_FEC.Data[2849] := 571.41;
   Prof_FEC.Data[2850] := 531.57;
   Prof_FEC.Data[2851] := 531.87;
   Prof_FEC.Data[2852] := 452.97;
   Prof_FEC.Data[2853] := 353.13;
   Prof_FEC.Data[2854] := 348.14;
   Prof_FEC.Data[2855] := 324.08;
   Prof_FEC.Data[2856] := 290.35;
   Prof_FEC.Data[2857] := 260.8;
   Prof_FEC.Data[2858] := 254.14;
   Prof_FEC.Data[2859] := 275.22;
   Prof_FEC.Data[2860] := 42.512;
   Prof_FEC.Data[2861] := 43.985;
   Prof_FEC.Data[2862] := 48.395;
   Prof_FEC.Data[2863] := 44.67;
   Prof_FEC.Data[2864] := 42.269;
   Prof_FEC.Data[2865] := 43.399;
   Prof_FEC.Data[2866] := 43.075;
   Prof_FEC.Data[2867] := 42.471;
   Prof_FEC.Data[2868] := 44.191;
   Prof_FEC.Data[2869] := 47.121;
   Prof_FEC.Data[2870] := 46.855;
   Prof_FEC.Data[2871] := 45.065;
   Prof_FEC.Data[2872] := 45.497;
   Prof_FEC.Data[2873] := 44.449;
   Prof_FEC.Data[2874] := 45.185;
   Prof_FEC.Data[2875] := 46.088;
   Prof_FEC.Data[2876] := 45.99;
   Prof_FEC.Data[2877] := 46.974;
   Prof_FEC.Data[2878] := 48.985;
   Prof_FEC.Data[2879] := 50.0;
   Prof_FEC.Data[2880] := 50.0;
   Prof_FEC.Data[2881] := 44.497;
   Prof_FEC.Data[2882] := 44.025;
   Prof_FEC.Data[2883] := 42.434;
   Prof_FEC.Data[2884] := 50.0;
   Prof_FEC.Data[2885] := 50.0;
   Prof_FEC.Data[2886] := 50.0;
   Prof_FEC.Data[2887] := 48.332;
   Prof_FEC.Data[2888] := 50.0;
   Prof_FEC.Data[2889] := 49.962;
   Prof_FEC.Data[2890] := 49.284;
   Prof_FEC.Data[2891] := 50.0;
   Prof_FEC.Data[2892] := 50.0;
   Prof_FEC.Data[2893] := 50.0;
   Prof_FEC.Data[2894] := 50.0;
   Prof_FEC.Data[2895] := 49.389;
   Prof_FEC.Data[2896] := 47.822;
   Prof_FEC.Data[2897] := 47.859;
   Prof_FEC.Data[2898] := 47.806;
   Prof_FEC.Data[2899] := 49.44;
   Prof_FEC.Data[2900] := 346.12;
   Prof_FEC.Data[2901] := 371.02;
   Prof_FEC.Data[2902] := 369.33;
   Prof_FEC.Data[2903] := 364.86;
   Prof_FEC.Data[2904] := 404.37;
   Prof_FEC.Data[2905] := 432.41;
   Prof_FEC.Data[2906] := 462.05;
   Prof_FEC.Data[2907] := 475.67;
   Prof_FEC.Data[2908] := 570.16;
   Prof_FEC.Data[2909] := 568.03;
   Prof_FEC.Data[2910] := 634.48;
   Prof_FEC.Data[2911] := 603.18;
   Prof_FEC.Data[2912] := 631.56;
   Prof_FEC.Data[2913] := 644.03;
   Prof_FEC.Data[2914] := 671.29;
   Prof_FEC.Data[2915] := 653.71;
   Prof_FEC.Data[2916] := 748.65;
   Prof_FEC.Data[2917] := 721.98;
   Prof_FEC.Data[2918] := 746.11;
   Prof_FEC.Data[2919] := 756.87;
   Prof_FEC.Data[2920] := 753.7;
   Prof_FEC.Data[2921] := 690.9;
   Prof_FEC.Data[2922] := 643.43;
   Prof_FEC.Data[2923] := 768.11;
   Prof_FEC.Data[2924] := 739.92;
   Prof_FEC.Data[2925] := 698.53;
   Prof_FEC.Data[2926] := 662.15;
   Prof_FEC.Data[2927] := 730.13;
   Prof_FEC.Data[2928] := 631.34;
   Prof_FEC.Data[2929] := 661.64;
   Prof_FEC.Data[2930] := 661.2;
   Prof_FEC.Data[2931] := 657.85;
   Prof_FEC.Data[2932] := 645.99;
   Prof_FEC.Data[2933] := 674.94;
   Prof_FEC.Data[2934] := 626.24;
   Prof_FEC.Data[2935] := 664.68;
   Prof_FEC.Data[2936] := 654.97;
   Prof_FEC.Data[2937] := 624.84;
   Prof_FEC.Data[2938] := 586.06;
   Prof_FEC.Data[2939] := 636.68;
   Prof_FEC.Data[2940] := 535.18;
   Prof_FEC.Data[2941] := 619.14;
   Prof_FEC.Data[2942] := 579.71;
   Prof_FEC.Data[2943] := 718.49;
   Prof_FEC.Data[2944] := 702.83;
   Prof_FEC.Data[2945] := 748.19;
   Prof_FEC.Data[2946] := 742.36;
   Prof_FEC.Data[2947] := 631.83;
   Prof_FEC.Data[2948] := 562.51;
   Prof_FEC.Data[2949] := 439.31;
   Prof_FEC.Data[2950] := 392.79;
   Prof_FEC.Data[2951] := 358.16;
   Prof_FEC.Data[2952] := 336.6;
   Prof_FEC.Data[2953] := 270.6;
   Prof_FEC.Data[2954] := 300.12;
   Prof_FEC.Data[2955] := 298.55;
   Prof_FEC.Data[2956] := 50.0;
   Prof_FEC.Data[2957] := 50.0;
   Prof_FEC.Data[2958] := 50.0;
   Prof_FEC.Data[2959] := 50.0;
   Prof_FEC.Data[2960] := 46.25;
   Prof_FEC.Data[2961] := 46.329;
   Prof_FEC.Data[2962] := 45.577;
   Prof_FEC.Data[2963] := 49.086;
   Prof_FEC.Data[2964] := 48.826;
   Prof_FEC.Data[2965] := 50.0;
   Prof_FEC.Data[2966] := 47.324;
   Prof_FEC.Data[2967] := 50.0;
   Prof_FEC.Data[2968] := 47.209;
   Prof_FEC.Data[2969] := 46.848;
   Prof_FEC.Data[2970] := 47.068;
   Prof_FEC.Data[2971] := 48.621;
   Prof_FEC.Data[2972] := 50.0;
   Prof_FEC.Data[2973] := 50.0;
   Prof_FEC.Data[2974] := 50.0;
   Prof_FEC.Data[2975] := 47.922;
   Prof_FEC.Data[2976] := 50.0;
   Prof_FEC.Data[2977] := 50.0;
   Prof_FEC.Data[2978] := 44.343;
   Prof_FEC.Data[2979] := 46.784;
   Prof_FEC.Data[2980] := 50.0;
   Prof_FEC.Data[2981] := 50.0;
   Prof_FEC.Data[2982] := 50.0;
   Prof_FEC.Data[2983] := 50.0;
   Prof_FEC.Data[2984] := 43.206;
   Prof_FEC.Data[2985] := 48.171;
   Prof_FEC.Data[2986] := 47.023;
   Prof_FEC.Data[2987] := 49.191;
   Prof_FEC.Data[2988] := 48.539;
   Prof_FEC.Data[2989] := 48.828;
   Prof_FEC.Data[2990] := 49.635;
   Prof_FEC.Data[2991] := 50.0;
   Prof_FEC.Data[2992] := 48.642;
   Prof_FEC.Data[2993] := 43.155;
   Prof_FEC.Data[2994] := 42.138;
   Prof_FEC.Data[2995] := 48.491;
   Prof_FEC.Data[2996] := 304.15;
   Prof_FEC.Data[2997] := 330.3;
   Prof_FEC.Data[2998] := 293.38;
   Prof_FEC.Data[2999] := 295.95;
   Prof_FEC.Data[3000] := 250.4;
   Prof_FEC.Data[3001] := 254.13;
   Prof_FEC.Data[3002] := 259.08;
   Prof_FEC.Data[3003] := 289.43;
   Prof_FEC.Data[3004] := 332.74;
   Prof_FEC.Data[3005] := 358.91;
   Prof_FEC.Data[3006] := 404.18;
   Prof_FEC.Data[3007] := 342.93;
   Prof_FEC.Data[3008] := 280.6;
   Prof_FEC.Data[3009] := 278.51;
   Prof_FEC.Data[3010] := 279.12;
   Prof_FEC.Data[3011] := 297.34;
   Prof_FEC.Data[3012] := 377.75;
   Prof_FEC.Data[3013] := 378.44;
   Prof_FEC.Data[3014] := 390.01;
   Prof_FEC.Data[3015] := 338.01;
   Prof_FEC.Data[3016] := 353.61;
   Prof_FEC.Data[3017] := 338.59;
   Prof_FEC.Data[3018] := 377.26;
   Prof_FEC.Data[3019] := 392.97;
   Prof_FEC.Data[3020] := 398.59;
   Prof_FEC.Data[3021] := 379.43;
   Prof_FEC.Data[3022] := 371.59;
   Prof_FEC.Data[3023] := 353.14;
   Prof_FEC.Data[3024] := 323.14;
   Prof_FEC.Data[3025] := 286.45;
   Prof_FEC.Data[3026] := 262.12;
   Prof_FEC.Data[3027] := 254.31;
   Prof_FEC.Data[3028] := 280.31;
   Prof_FEC.Data[3029] := 281.23;
   Prof_FEC.Data[3030] := 286.18;
   Prof_FEC.Data[3031] := 289.28;
   Prof_FEC.Data[3032] := 314.49;
   Prof_FEC.Data[3033] := 312.86;
   Prof_FEC.Data[3034] := 287.4;
   Prof_FEC.Data[3035] := 254.42;
   Prof_FEC.Data[3036] := 337.05;
   Prof_FEC.Data[3037] := 317.9;
   Prof_FEC.Data[3038] := 292.07;
   Prof_FEC.Data[3039] := 273.2;
   Prof_FEC.Data[3040] := 207.56;
   Prof_FEC.Data[3041] := 175.2;
   Prof_FEC.Data[3042] := 163.44;
   Prof_FEC.Data[3043] := 215.63;
   Prof_FEC.Data[3044] := 234.15;
   Prof_FEC.Data[3045] := 250.68;
   Prof_FEC.Data[3046] := 269.4;
   Prof_FEC.Data[3047] := 266.43;
   Prof_FEC.Data[3048] := 282.15;
   Prof_FEC.Data[3049] := 292.66;
   Prof_FEC.Data[3050] := 275.18;
   Prof_FEC.Data[3051] := 277.22;
   Prof_FEC.Data[3052] := 41.715;
   Prof_FEC.Data[3053] := 39.062;
   Prof_FEC.Data[3054] := 42.719;
   Prof_FEC.Data[3055] := 42.928;
   Prof_FEC.Data[3056] := 47.383;
   Prof_FEC.Data[3057] := 44.237;
   Prof_FEC.Data[3058] := 47.256;
   Prof_FEC.Data[3059] := 44.542;
   Prof_FEC.Data[3060] := 43.998;
   Prof_FEC.Data[3061] := 45.672;
   Prof_FEC.Data[3062] := 42.611;
   Prof_FEC.Data[3063] := 47.856;
   Prof_FEC.Data[3064] := 48.829;
   Prof_FEC.Data[3065] := 47.605;
   Prof_FEC.Data[3066] := 50.0;
   Prof_FEC.Data[3067] := 47.645;
   Prof_FEC.Data[3068] := 45.197;
   Prof_FEC.Data[3069] := 43.021;
   Prof_FEC.Data[3070] := 42.577;
   Prof_FEC.Data[3071] := 43.107;
   Prof_FEC.Data[3072] := 46.925;
   Prof_FEC.Data[3073] := 47.577;
   Prof_FEC.Data[3074] := 41.953;
   Prof_FEC.Data[3075] := 43.543;
   Prof_FEC.Data[3076] := 40.381;
   Prof_FEC.Data[3077] := 38.77;
   Prof_FEC.Data[3078] := 41.083;
   Prof_FEC.Data[3079] := 43.29;
   Prof_FEC.Data[3080] := 47.103;
   Prof_FEC.Data[3081] := 49.23;
   Prof_FEC.Data[3082] := 50.0;
   Prof_FEC.Data[3083] := 46.789;
   Prof_FEC.Data[3084] := 48.025;
   Prof_FEC.Data[3085] := 43.33;
   Prof_FEC.Data[3086] := 41.971;
   Prof_FEC.Data[3087] := 46.349;
   Prof_FEC.Data[3088] := 50.0;
   Prof_FEC.Data[3089] := 45.259;
   Prof_FEC.Data[3090] := 50.0;
   Prof_FEC.Data[3091] := 47.031;
   Prof_FEC.Data[3092] := 280.25;
   Prof_FEC.Data[3093] := 275.08;
   Prof_FEC.Data[3094] := 302.18;
   Prof_FEC.Data[3095] := 322.06;
   Prof_FEC.Data[3096] := 331.52;
   Prof_FEC.Data[3097] := 316.81;
   Prof_FEC.Data[3098] := 338.58;
   Prof_FEC.Data[3099] := 323.82;
   Prof_FEC.Data[3100] := 291.16;
   Prof_FEC.Data[3101] := 258.55;
   Prof_FEC.Data[3102] := 259.35;
   Prof_FEC.Data[3103] := 242.41;
   Prof_FEC.Data[3104] := 250.48;
   Prof_FEC.Data[3105] := 253.94;
   Prof_FEC.Data[3106] := 232.93;
   Prof_FEC.Data[3107] := 220.14;
   Prof_FEC.Data[3108] := 200.41;
   Prof_FEC.Data[3109] := 180.8;
   Prof_FEC.Data[3110] := 160.44;
   Prof_FEC.Data[3111] := 186.66;
   Prof_FEC.Data[3112] := 195.2;
   Prof_FEC.Data[3113] := 234.93;
   Prof_FEC.Data[3114] := 189.38;
   Prof_FEC.Data[3115] := 191.48;
   Prof_FEC.Data[3116] := 180.23;
   Prof_FEC.Data[3117] := 159.63;
   Prof_FEC.Data[3118] := 137.94;
   Prof_FEC.Data[3119] := 151.78;
   Prof_FEC.Data[3120] := 181.73;
   Prof_FEC.Data[3121] := 191.55;
   Prof_FEC.Data[3122] := 199.23;
   Prof_FEC.Data[3123] := 200.33;
   Prof_FEC.Data[3124] := 155.06;
   Prof_FEC.Data[3125] := 175.09;
   Prof_FEC.Data[3126] := 152.74;
   Prof_FEC.Data[3127] := 160.0;
   Prof_FEC.Data[3128] := 195.68;
   Prof_FEC.Data[3129] := 186.25;
   Prof_FEC.Data[3130] := 204.27;
   Prof_FEC.Data[3131] := 193.14;
   Prof_FEC.Data[3132] := 161.76;
   Prof_FEC.Data[3133] := 166.2;
   Prof_FEC.Data[3134] := 155.86;
   Prof_FEC.Data[3135] := 167.93;
   Prof_FEC.Data[3136] := 167.48;
   Prof_FEC.Data[3137] := 201.59;
   Prof_FEC.Data[3138] := 196.02;
   Prof_FEC.Data[3139] := 224.77;
   Prof_FEC.Data[3140] := 281.19;
   Prof_FEC.Data[3141] := 271.62;
   Prof_FEC.Data[3142] := 309.48;
   Prof_FEC.Data[3143] := 310.68;
   Prof_FEC.Data[3144] := 297.31;
   Prof_FEC.Data[3145] := 309.21;
   Prof_FEC.Data[3146] := 308.46;
   Prof_FEC.Data[3147] := 311.34;
   Prof_FEC.Data[3148] := 43.62;
   Prof_FEC.Data[3149] := 42.745;
   Prof_FEC.Data[3150] := 39.66;
   Prof_FEC.Data[3151] := 44.482;
   Prof_FEC.Data[3152] := 49.469;
   Prof_FEC.Data[3153] := 50.0;
   Prof_FEC.Data[3154] := 49.925;
   Prof_FEC.Data[3155] := 50.0;
   Prof_FEC.Data[3156] := 45.695;
   Prof_FEC.Data[3157] := 45.073;
   Prof_FEC.Data[3158] := 45.69;
   Prof_FEC.Data[3159] := 47.916;
   Prof_FEC.Data[3160] := 49.692;
   Prof_FEC.Data[3161] := 50.0;
   Prof_FEC.Data[3162] := 50.0;
   Prof_FEC.Data[3163] := 49.179;
   Prof_FEC.Data[3164] := 49.953;
   Prof_FEC.Data[3165] := 47.408;
   Prof_FEC.Data[3166] := 47.211;
   Prof_FEC.Data[3167] := 46.58;
   Prof_FEC.Data[3168] := 50.0;
   Prof_FEC.Data[3169] := 50.0;
   Prof_FEC.Data[3170] := 50.0;
   Prof_FEC.Data[3171] := 50.0;
   Prof_FEC.Data[3172] := 46.857;
   Prof_FEC.Data[3173] := 45.372;
   Prof_FEC.Data[3174] := 47.685;
   Prof_FEC.Data[3175] := 46.23;
   Prof_FEC.Data[3176] := 50.0;
   Prof_FEC.Data[3177] := 48.176;
   Prof_FEC.Data[3178] := 49.865;
   Prof_FEC.Data[3179] := 50.0;
   Prof_FEC.Data[3180] := 49.463;
   Prof_FEC.Data[3181] := 47.717;
   Prof_FEC.Data[3182] := 46.007;
   Prof_FEC.Data[3183] := 45.044;
   Prof_FEC.Data[3184] := 50.0;
   Prof_FEC.Data[3185] := 49.21;
   Prof_FEC.Data[3186] := 50.0;
   Prof_FEC.Data[3187] := 49.134;
   Prof_FEC.Data[3188] := 346.39;
   Prof_FEC.Data[3189] := 289.36;
   Prof_FEC.Data[3190] := 333.52;
   Prof_FEC.Data[3191] := 317.49;
   Prof_FEC.Data[3192] := 369.82;
   Prof_FEC.Data[3193] := 383.47;
   Prof_FEC.Data[3194] := 415.51;
   Prof_FEC.Data[3195] := 443.19;
   Prof_FEC.Data[3196] := 467.72;
   Prof_FEC.Data[3197] := 497.05;
   Prof_FEC.Data[3198] := 477.64;
   Prof_FEC.Data[3199] := 519.41;
   Prof_FEC.Data[3200] := 475.47;
   Prof_FEC.Data[3201] := 544.8;
   Prof_FEC.Data[3202] := 554.14;
   Prof_FEC.Data[3203] := 607.38;
   Prof_FEC.Data[3204] := 601.27;
   Prof_FEC.Data[3205] := 646.27;
   Prof_FEC.Data[3206] := 621.28;
   Prof_FEC.Data[3207] := 575.74;
   Prof_FEC.Data[3208] := 654.1;
   Prof_FEC.Data[3209] := 666.23;
   Prof_FEC.Data[3210] := 658.97;
   Prof_FEC.Data[3211] := 728.59;
   Prof_FEC.Data[3212] := 616.05;
   Prof_FEC.Data[3213] := 700.7;
   Prof_FEC.Data[3214] := 694.08;
   Prof_FEC.Data[3215] := 640.1;
   Prof_FEC.Data[3216] := 632.22;
   Prof_FEC.Data[3217] := 647.57;
   Prof_FEC.Data[3218] := 630.77;
   Prof_FEC.Data[3219] := 645.02;
   Prof_FEC.Data[3220] := 681.65;
   Prof_FEC.Data[3221] := 666.04;
   Prof_FEC.Data[3222] := 728.09;
   Prof_FEC.Data[3223] := 730.62;
   Prof_FEC.Data[3224] := 696.56;
   Prof_FEC.Data[3225] := 717.1;
   Prof_FEC.Data[3226] := 732.7;
   Prof_FEC.Data[3227] := 774.81;
   Prof_FEC.Data[3228] := 723.82;
   Prof_FEC.Data[3229] := 636.53;
   Prof_FEC.Data[3230] := 645.48;
   Prof_FEC.Data[3231] := 700.3;
   Prof_FEC.Data[3232] := 698.29;
   Prof_FEC.Data[3233] := 737.81;
   Prof_FEC.Data[3234] := 759.11;
   Prof_FEC.Data[3235] := 662.35;
   Prof_FEC.Data[3236] := 477.19;
   Prof_FEC.Data[3237] := 481.71;
   Prof_FEC.Data[3238] := 390.5;
   Prof_FEC.Data[3239] := 377.19;
   Prof_FEC.Data[3240] := 333.67;
   Prof_FEC.Data[3241] := 309.25;
   Prof_FEC.Data[3242] := 280.6;
   Prof_FEC.Data[3243] := 262.0;
   Prof_FEC.Data[3244] := 46.074;
   Prof_FEC.Data[3245] := 45.026;
   Prof_FEC.Data[3246] := 49.148;
   Prof_FEC.Data[3247] := 48.0;
   Prof_FEC.Data[3248] := 44.833;
   Prof_FEC.Data[3249] := 42.146;
   Prof_FEC.Data[3250] := 44.026;
   Prof_FEC.Data[3251] := 46.4;
   Prof_FEC.Data[3252] := 47.411;
   Prof_FEC.Data[3253] := 50.0;
   Prof_FEC.Data[3254] := 48.055;
   Prof_FEC.Data[3255] := 46.331;
   Prof_FEC.Data[3256] := 42.053;
   Prof_FEC.Data[3257] := 44.033;
   Prof_FEC.Data[3258] := 42.903;
   Prof_FEC.Data[3259] := 41.375;
   Prof_FEC.Data[3260] := 43.489;
   Prof_FEC.Data[3261] := 42.959;
   Prof_FEC.Data[3262] := 41.619;
   Prof_FEC.Data[3263] := 38.252;
   Prof_FEC.Data[3264] := 39.143;
   Prof_FEC.Data[3265] := 44.39;
   Prof_FEC.Data[3266] := 43.997;
   Prof_FEC.Data[3267] := 44.809;
   Prof_FEC.Data[3268] := 44.855;
   Prof_FEC.Data[3269] := 49.874;
   Prof_FEC.Data[3270] := 49.062;
   Prof_FEC.Data[3271] := 49.984;
   Prof_FEC.Data[3272] := 44.153;
   Prof_FEC.Data[3273] := 44.051;
   Prof_FEC.Data[3274] := 45.474;
   Prof_FEC.Data[3275] := 48.575;
   Prof_FEC.Data[3276] := 47.434;
   Prof_FEC.Data[3277] := 47.226;
   Prof_FEC.Data[3278] := 50.0;
   Prof_FEC.Data[3279] := 44.289;
   Prof_FEC.Data[3280] := 43.117;
   Prof_FEC.Data[3281] := 44.671;
   Prof_FEC.Data[3282] := 46.71;
   Prof_FEC.Data[3283] := 44.17;
   Prof_FEC.Data[3284] := 310.65;
   Prof_FEC.Data[3285] := 314.78;
   Prof_FEC.Data[3286] := 329.04;
   Prof_FEC.Data[3287] := 312.36;
   Prof_FEC.Data[3288] := 364.24;
   Prof_FEC.Data[3289] := 367.32;
   Prof_FEC.Data[3290] := 406.77;
   Prof_FEC.Data[3291] := 423.93;
   Prof_FEC.Data[3292] := 487.1;
   Prof_FEC.Data[3293] := 475.59;
   Prof_FEC.Data[3294] := 474.24;
   Prof_FEC.Data[3295] := 596.67;
   Prof_FEC.Data[3296] := 495.72;
   Prof_FEC.Data[3297] := 526.67;
   Prof_FEC.Data[3298] := 554.68;
   Prof_FEC.Data[3299] := 611.85;
   Prof_FEC.Data[3300] := 630.65;
   Prof_FEC.Data[3301] := 697.53;
   Prof_FEC.Data[3302] := 752.38;
   Prof_FEC.Data[3303] := 781.49;
   Prof_FEC.Data[3304] := 689.8;
   Prof_FEC.Data[3305] := 673.84;
   Prof_FEC.Data[3306] := 615.77;
   Prof_FEC.Data[3307] := 690.63;
   Prof_FEC.Data[3308] := 684.53;
   Prof_FEC.Data[3309] := 577.83;
   Prof_FEC.Data[3310] := 601.23;
   Prof_FEC.Data[3311] := 676.74;
   Prof_FEC.Data[3312] := 621.85;
   Prof_FEC.Data[3313] := 582.04;
   Prof_FEC.Data[3314] := 581.97;
   Prof_FEC.Data[3315] := 604.97;
   Prof_FEC.Data[3316] := 666.68;
   Prof_FEC.Data[3317] := 668.5;
   Prof_FEC.Data[3318] := 684.96;
   Prof_FEC.Data[3319] := 604.3;
   Prof_FEC.Data[3320] := 562.65;
   Prof_FEC.Data[3321] := 561.05;
   Prof_FEC.Data[3322] := 611.11;
   Prof_FEC.Data[3323] := 631.0;
   Prof_FEC.Data[3324] := 631.94;
   Prof_FEC.Data[3325] := 658.22;
   Prof_FEC.Data[3326] := 710.56;
   Prof_FEC.Data[3327] := 695.95;
   Prof_FEC.Data[3328] := 754.97;
   Prof_FEC.Data[3329] := 777.82;
   Prof_FEC.Data[3330] := 698.01;
   Prof_FEC.Data[3331] := 591.61;
   Prof_FEC.Data[3332] := 492.29;
   Prof_FEC.Data[3333] := 457.9;
   Prof_FEC.Data[3334] := 404.33;
   Prof_FEC.Data[3335] := 337.98;
   Prof_FEC.Data[3336] := 317.57;
   Prof_FEC.Data[3337] := 251.71;
   Prof_FEC.Data[3338] := 234.37;
   Prof_FEC.Data[3339] := 235.24;
   Prof_FEC.Data[3340] := 43.505;
   Prof_FEC.Data[3341] := 47.144;
   Prof_FEC.Data[3342] := 45.247;
   Prof_FEC.Data[3343] := 45.176;
   Prof_FEC.Data[3344] := 41.617;
   Prof_FEC.Data[3345] := 41.578;
   Prof_FEC.Data[3346] := 41.097;
   Prof_FEC.Data[3347] := 42.725;
   Prof_FEC.Data[3348] := 41.475;
   Prof_FEC.Data[3349] := 44.21;
   Prof_FEC.Data[3350] := 45.984;
   Prof_FEC.Data[3351] := 43.104;
   Prof_FEC.Data[3352] := 43.896;
   Prof_FEC.Data[3353] := 45.131;
   Prof_FEC.Data[3354] := 46.161;
   Prof_FEC.Data[3355] := 44.585;
   Prof_FEC.Data[3356] := 48.737;
   Prof_FEC.Data[3357] := 45.879;
   Prof_FEC.Data[3358] := 47.95;
   Prof_FEC.Data[3359] := 48.248;
   Prof_FEC.Data[3360] := 46.747;
   Prof_FEC.Data[3361] := 45.383;
   Prof_FEC.Data[3362] := 43.62;
   Prof_FEC.Data[3363] := 45.106;
   Prof_FEC.Data[3364] := 50.0;
   Prof_FEC.Data[3365] := 50.0;
   Prof_FEC.Data[3366] := 50.0;
   Prof_FEC.Data[3367] := 50.0;
   Prof_FEC.Data[3368] := 49.23;
   Prof_FEC.Data[3369] := 44.168;
   Prof_FEC.Data[3370] := 46.647;
   Prof_FEC.Data[3371] := 47.707;
   Prof_FEC.Data[3372] := 50.0;
   Prof_FEC.Data[3373] := 50.0;
   Prof_FEC.Data[3374] := 50.0;
   Prof_FEC.Data[3375] := 50.0;
   Prof_FEC.Data[3376] := 49.503;
   Prof_FEC.Data[3377] := 50.0;
   Prof_FEC.Data[3378] := 50.0;
   Prof_FEC.Data[3379] := 50.0;
   Prof_FEC.Data[3380] := 358.32;
   Prof_FEC.Data[3381] := 405.51;
   Prof_FEC.Data[3382] := 397.33;
   Prof_FEC.Data[3383] := 431.99;
   Prof_FEC.Data[3384] := 430.28;
   Prof_FEC.Data[3385] := 477.66;
   Prof_FEC.Data[3386] := 476.1;
   Prof_FEC.Data[3387] := 489.56;
   Prof_FEC.Data[3388] := 509.03;
   Prof_FEC.Data[3389] := 532.7;
   Prof_FEC.Data[3390] := 562.67;
   Prof_FEC.Data[3391] := 586.62;
   Prof_FEC.Data[3392] := 562.96;
   Prof_FEC.Data[3393] := 593.98;
   Prof_FEC.Data[3394] := 694.87;
   Prof_FEC.Data[3395] := 643.68;
   Prof_FEC.Data[3396] := 699.75;
   Prof_FEC.Data[3397] := 699.41;
   Prof_FEC.Data[3398] := 740.64;
   Prof_FEC.Data[3399] := 755.2;
   Prof_FEC.Data[3400] := 677.01;
   Prof_FEC.Data[3401] := 749.41;
   Prof_FEC.Data[3402] := 792.63;
   Prof_FEC.Data[3403] := 693.04;
   Prof_FEC.Data[3404] := 649.7;
   Prof_FEC.Data[3405] := 722.86;
   Prof_FEC.Data[3406] := 648.54;
   Prof_FEC.Data[3407] := 704.1;
   Prof_FEC.Data[3408] := 598.06;
   Prof_FEC.Data[3409] := 674.99;
   Prof_FEC.Data[3410] := 601.34;
   Prof_FEC.Data[3411] := 627.49;
   Prof_FEC.Data[3412] := 569.41;
   Prof_FEC.Data[3413] := 631.76;
   Prof_FEC.Data[3414] := 608.13;
   Prof_FEC.Data[3415] := 609.53;
   Prof_FEC.Data[3416] := 666.17;
   Prof_FEC.Data[3417] := 596.03;
   Prof_FEC.Data[3418] := 636.34;
   Prof_FEC.Data[3419] := 642.26;
   Prof_FEC.Data[3420] := 709.47;
   Prof_FEC.Data[3421] := 702.28;
   Prof_FEC.Data[3422] := 692.44;
   Prof_FEC.Data[3423] := 623.9;
   Prof_FEC.Data[3424] := 754.27;
   Prof_FEC.Data[3425] := 676.35;
   Prof_FEC.Data[3426] := 627.92;
   Prof_FEC.Data[3427] := 562.01;
   Prof_FEC.Data[3428] := 470.7;
   Prof_FEC.Data[3429] := 424.42;
   Prof_FEC.Data[3430] := 374.66;
   Prof_FEC.Data[3431] := 372.53;
   Prof_FEC.Data[3432] := 294.12;
   Prof_FEC.Data[3433] := 322.82;
   Prof_FEC.Data[3434] := 301.32;
   Prof_FEC.Data[3435] := 307.34;
   Prof_FEC.Data[3436] := 48.963;
   Prof_FEC.Data[3437] := 50.0;
   Prof_FEC.Data[3438] := 50.0;
   Prof_FEC.Data[3439] := 48.131;
   Prof_FEC.Data[3440] := 44.201;
   Prof_FEC.Data[3441] := 45.255;
   Prof_FEC.Data[3442] := 46.306;
   Prof_FEC.Data[3443] := 44.405;
   Prof_FEC.Data[3444] := 45.955;
   Prof_FEC.Data[3445] := 48.734;
   Prof_FEC.Data[3446] := 50.0;
   Prof_FEC.Data[3447] := 50.0;
   Prof_FEC.Data[3448] := 46.932;
   Prof_FEC.Data[3449] := 45.854;
   Prof_FEC.Data[3450] := 47.503;
   Prof_FEC.Data[3451] := 46.317;
   Prof_FEC.Data[3452] := 50.0;
   Prof_FEC.Data[3453] := 50.0;
   Prof_FEC.Data[3454] := 50.0;
   Prof_FEC.Data[3455] := 50.0;
   Prof_FEC.Data[3456] := 50.0;
   Prof_FEC.Data[3457] := 46.162;
   Prof_FEC.Data[3458] := 49.522;
   Prof_FEC.Data[3459] := 50.0;
   Prof_FEC.Data[3460] := 50.0;
   Prof_FEC.Data[3461] := 50.0;
   Prof_FEC.Data[3462] := 47.872;
   Prof_FEC.Data[3463] := 48.82;
   Prof_FEC.Data[3464] := 46.15;
   Prof_FEC.Data[3465] := 49.967;
   Prof_FEC.Data[3466] := 46.093;
   Prof_FEC.Data[3467] := 46.895;
   Prof_FEC.Data[3468] := 49.285;
   Prof_FEC.Data[3469] := 50.0;
   Prof_FEC.Data[3470] := 50.0;
   Prof_FEC.Data[3471] := 44.015;
   Prof_FEC.Data[3472] := 45.429;
   Prof_FEC.Data[3473] := 45.914;
   Prof_FEC.Data[3474] := 48.1;
   Prof_FEC.Data[3475] := 45.012;
   Prof_FEC.Data[3476] := 328.14;
   Prof_FEC.Data[3477] := 329.73;
   Prof_FEC.Data[3478] := 388.89;
   Prof_FEC.Data[3479] := 386.52;
   Prof_FEC.Data[3480] := 380.63;
   Prof_FEC.Data[3481] := 438.4;
   Prof_FEC.Data[3482] := 448.93;
   Prof_FEC.Data[3483] := 475.18;
   Prof_FEC.Data[3484] := 482.55;
   Prof_FEC.Data[3485] := 523.9;
   Prof_FEC.Data[3486] := 544.34;
   Prof_FEC.Data[3487] := 620.31;
   Prof_FEC.Data[3488] := 552.31;
   Prof_FEC.Data[3489] := 560.55;
   Prof_FEC.Data[3490] := 614.8;
   Prof_FEC.Data[3491] := 673.81;
   Prof_FEC.Data[3492] := 646.93;
   Prof_FEC.Data[3493] := 705.29;
   Prof_FEC.Data[3494] := 665.37;
   Prof_FEC.Data[3495] := 739.15;
   Prof_FEC.Data[3496] := 695.2;
   Prof_FEC.Data[3497] := 772.17;
   Prof_FEC.Data[3498] := 778.09;
   Prof_FEC.Data[3499] := 723.9;
   Prof_FEC.Data[3500] := 744.61;
   Prof_FEC.Data[3501] := 728.83;
   Prof_FEC.Data[3502] := 709.02;
   Prof_FEC.Data[3503] := 693.02;
   Prof_FEC.Data[3504] := 657.92;
   Prof_FEC.Data[3505] := 634.33;
   Prof_FEC.Data[3506] := 650.7;
   Prof_FEC.Data[3507] := 611.98;
   Prof_FEC.Data[3508] := 682.67;
   Prof_FEC.Data[3509] := 668.64;
   Prof_FEC.Data[3510] := 705.81;
   Prof_FEC.Data[3511] := 748.53;
   Prof_FEC.Data[3512] := 686.13;
   Prof_FEC.Data[3513] := 609.32;
   Prof_FEC.Data[3514] := 668.24;
   Prof_FEC.Data[3515] := 704.27;
   Prof_FEC.Data[3516] := 666.28;
   Prof_FEC.Data[3517] := 694.74;
   Prof_FEC.Data[3518] := 617.53;
   Prof_FEC.Data[3519] := 646.54;
   Prof_FEC.Data[3520] := 710.56;
   Prof_FEC.Data[3521] := 745.57;
   Prof_FEC.Data[3522] := 670.89;
   Prof_FEC.Data[3523] := 678.75;
   Prof_FEC.Data[3524] := 559.3;
   Prof_FEC.Data[3525] := 445.37;
   Prof_FEC.Data[3526] := 432.65;
   Prof_FEC.Data[3527] := 366.26;
   Prof_FEC.Data[3528] := 334.74;
   Prof_FEC.Data[3529] := 306.28;
   Prof_FEC.Data[3530] := 310.24;
   Prof_FEC.Data[3531] := 322.86;
   Prof_FEC.Data[3532] := 50.0;
   Prof_FEC.Data[3533] := 50.0;
   Prof_FEC.Data[3534] := 50.0;
   Prof_FEC.Data[3535] := 49.405;
   Prof_FEC.Data[3536] := 49.783;
   Prof_FEC.Data[3537] := 42.422;
   Prof_FEC.Data[3538] := 48.392;
   Prof_FEC.Data[3539] := 48.286;
   Prof_FEC.Data[3540] := 50.0;
   Prof_FEC.Data[3541] := 50.0;
   Prof_FEC.Data[3542] := 47.503;
   Prof_FEC.Data[3543] := 49.875;
   Prof_FEC.Data[3544] := 45.983;
   Prof_FEC.Data[3545] := 45.691;
   Prof_FEC.Data[3546] := 44.153;
   Prof_FEC.Data[3547] := 47.806;
   Prof_FEC.Data[3548] := 49.91;
   Prof_FEC.Data[3549] := 49.475;
   Prof_FEC.Data[3550] := 49.494;
   Prof_FEC.Data[3551] := 45.933;
   Prof_FEC.Data[3552] := 43.953;
   Prof_FEC.Data[3553] := 44.087;
   Prof_FEC.Data[3554] := 45.228;
   Prof_FEC.Data[3555] := 46.511;
   Prof_FEC.Data[3556] := 50.0;
   Prof_FEC.Data[3557] := 50.0;
   Prof_FEC.Data[3558] := 49.666;
   Prof_FEC.Data[3559] := 48.395;
   Prof_FEC.Data[3560] := 47.539;
   Prof_FEC.Data[3561] := 43.214;
   Prof_FEC.Data[3562] := 43.735;
   Prof_FEC.Data[3563] := 44.802;
   Prof_FEC.Data[3564] := 45.855;
   Prof_FEC.Data[3565] := 46.384;
   Prof_FEC.Data[3566] := 46.643;
   Prof_FEC.Data[3567] := 49.813;
   Prof_FEC.Data[3568] := 44.822;
   Prof_FEC.Data[3569] := 41.242;
   Prof_FEC.Data[3570] := 42.94;
   Prof_FEC.Data[3571] := 42.81;
   Prof_FEC.Data[3572] := 280.52;
   Prof_FEC.Data[3573] := 280.78;
   Prof_FEC.Data[3574] := 308.35;
   Prof_FEC.Data[3575] := 272.47;
   Prof_FEC.Data[3576] := 285.11;
   Prof_FEC.Data[3577] := 329.03;
   Prof_FEC.Data[3578] := 327.23;
   Prof_FEC.Data[3579] := 412.59;
   Prof_FEC.Data[3580] := 385.62;
   Prof_FEC.Data[3581] := 408.94;
   Prof_FEC.Data[3582] := 471.82;
   Prof_FEC.Data[3583] := 423.37;
   Prof_FEC.Data[3584] := 487.71;
   Prof_FEC.Data[3585] := 511.75;
   Prof_FEC.Data[3586] := 568.7;
   Prof_FEC.Data[3587] := 562.85;
   Prof_FEC.Data[3588] := 628.31;
   Prof_FEC.Data[3589] := 625.45;
   Prof_FEC.Data[3590] := 672.82;
   Prof_FEC.Data[3591] := 658.03;
   Prof_FEC.Data[3592] := 685.68;
   Prof_FEC.Data[3593] := 721.75;
   Prof_FEC.Data[3594] := 655.04;
   Prof_FEC.Data[3595] := 675.8;
   Prof_FEC.Data[3596] := 758.5;
   Prof_FEC.Data[3597] := 672.75;
   Prof_FEC.Data[3598] := 595.17;
   Prof_FEC.Data[3599] := 649.49;
   Prof_FEC.Data[3600] := 576.06;
   Prof_FEC.Data[3601] := 652.64;
   Prof_FEC.Data[3602] := 662.64;
   Prof_FEC.Data[3603] := 725.24;
   Prof_FEC.Data[3604] := 767.6;
   Prof_FEC.Data[3605] := 774.92;
   Prof_FEC.Data[3606] := 678.79;
   Prof_FEC.Data[3607] := 693.24;
   Prof_FEC.Data[3608] := 719.53;
   Prof_FEC.Data[3609] := 613.5;
   Prof_FEC.Data[3610] := 631.46;
   Prof_FEC.Data[3611] := 653.44;
   Prof_FEC.Data[3612] := 658.91;
   Prof_FEC.Data[3613] := 673.06;
   Prof_FEC.Data[3614] := 643.05;
   Prof_FEC.Data[3615] := 666.58;
   Prof_FEC.Data[3616] := 690.83;
   Prof_FEC.Data[3617] := 709.93;
   Prof_FEC.Data[3618] := 643.17;
   Prof_FEC.Data[3619] := 579.0;
   Prof_FEC.Data[3620] := 521.64;
   Prof_FEC.Data[3621] := 429.37;
   Prof_FEC.Data[3622] := 406.69;
   Prof_FEC.Data[3623] := 342.36;
   Prof_FEC.Data[3624] := 345.78;
   Prof_FEC.Data[3625] := 313.28;
   Prof_FEC.Data[3626] := 274.87;
   Prof_FEC.Data[3627] := 297.06;
   Prof_FEC.Data[3628] := 48.681;
   Prof_FEC.Data[3629] := 50.0;
   Prof_FEC.Data[3630] := 50.0;
   Prof_FEC.Data[3631] := 46.669;
   Prof_FEC.Data[3632] := 41.107;
   Prof_FEC.Data[3633] := 46.507;
   Prof_FEC.Data[3634] := 45.959;
   Prof_FEC.Data[3635] := 46.764;
   Prof_FEC.Data[3636] := 49.554;
   Prof_FEC.Data[3637] := 49.384;
   Prof_FEC.Data[3638] := 48.555;
   Prof_FEC.Data[3639] := 48.485;
   Prof_FEC.Data[3640] := 46.463;
   Prof_FEC.Data[3641] := 47.695;
   Prof_FEC.Data[3642] := 47.977;
   Prof_FEC.Data[3643] := 46.864;
   Prof_FEC.Data[3644] := 49.039;
   Prof_FEC.Data[3645] := 50.0;
   Prof_FEC.Data[3646] := 47.963;
   Prof_FEC.Data[3647] := 50.0;
   Prof_FEC.Data[3648] := 47.144;
   Prof_FEC.Data[3649] := 45.889;
   Prof_FEC.Data[3650] := 42.252;
   Prof_FEC.Data[3651] := 45.608;
   Prof_FEC.Data[3652] := 46.753;
   Prof_FEC.Data[3653] := 47.297;
   Prof_FEC.Data[3654] := 46.02;
   Prof_FEC.Data[3655] := 47.015;
   Prof_FEC.Data[3656] := 44.139;
   Prof_FEC.Data[3657] := 44.546;
   Prof_FEC.Data[3658] := 41.938;
   Prof_FEC.Data[3659] := 38.349;
   Prof_FEC.Data[3660] := 45.583;
   Prof_FEC.Data[3661] := 42.694;
   Prof_FEC.Data[3662] := 43.026;
   Prof_FEC.Data[3663] := 45.724;
   Prof_FEC.Data[3664] := 41.133;
   Prof_FEC.Data[3665] := 44.281;
   Prof_FEC.Data[3666] := 42.76;
   Prof_FEC.Data[3667] := 44.791;
   Prof_FEC.Data[3668] := 312.73;
   Prof_FEC.Data[3669] := 358.53;
   Prof_FEC.Data[3670] := 346.07;
   Prof_FEC.Data[3671] := 312.08;
   Prof_FEC.Data[3672] := 329.21;
   Prof_FEC.Data[3673] := 273.82;
   Prof_FEC.Data[3674] := 296.46;
   Prof_FEC.Data[3675] := 282.57;
   Prof_FEC.Data[3676] := 313.57;
   Prof_FEC.Data[3677] := 313.71;
   Prof_FEC.Data[3678] := 318.99;
   Prof_FEC.Data[3679] := 320.61;
   Prof_FEC.Data[3680] := 275.51;
   Prof_FEC.Data[3681] := 285.15;
   Prof_FEC.Data[3682] := 286.08;
   Prof_FEC.Data[3683] := 339.73;
   Prof_FEC.Data[3684] := 362.84;
   Prof_FEC.Data[3685] := 410.42;
   Prof_FEC.Data[3686] := 374.74;
   Prof_FEC.Data[3687] := 380.03;
   Prof_FEC.Data[3688] := 433.14;
   Prof_FEC.Data[3689] := 471.32;
   Prof_FEC.Data[3690] := 483.61;
   Prof_FEC.Data[3691] := 428.06;
   Prof_FEC.Data[3692] := 424.48;
   Prof_FEC.Data[3693] := 435.79;
   Prof_FEC.Data[3694] := 400.17;
   Prof_FEC.Data[3695] := 381.17;
   Prof_FEC.Data[3696] := 342.47;
   Prof_FEC.Data[3697] := 347.91;
   Prof_FEC.Data[3698] := 323.44;
   Prof_FEC.Data[3699] := 335.78;
   Prof_FEC.Data[3700] := 291.24;
   Prof_FEC.Data[3701] := 323.67;
   Prof_FEC.Data[3702] := 303.04;
   Prof_FEC.Data[3703] := 344.17;
   Prof_FEC.Data[3704] := 322.39;
   Prof_FEC.Data[3705] := 307.3;
   Prof_FEC.Data[3706] := 288.43;
   Prof_FEC.Data[3707] := 297.63;
   Prof_FEC.Data[3708] := 320.44;
   Prof_FEC.Data[3709] := 337.94;
   Prof_FEC.Data[3710] := 319.49;
   Prof_FEC.Data[3711] := 298.3;
   Prof_FEC.Data[3712] := 214.33;
   Prof_FEC.Data[3713] := 164.98;
   Prof_FEC.Data[3714] := 174.85;
   Prof_FEC.Data[3715] := 198.83;
   Prof_FEC.Data[3716] := 244.19;
   Prof_FEC.Data[3717] := 282.59;
   Prof_FEC.Data[3718] := 296.38;
   Prof_FEC.Data[3719] := 288.06;
   Prof_FEC.Data[3720] := 301.93;
   Prof_FEC.Data[3721] := 314.04;
   Prof_FEC.Data[3722] := 298.04;
   Prof_FEC.Data[3723] := 285.48;
   Prof_FEC.Data[3724] := 39.69;
   Prof_FEC.Data[3725] := 42.335;
   Prof_FEC.Data[3726] := 45.25;
   Prof_FEC.Data[3727] := 44.971;
   Prof_FEC.Data[3728] := 47.55;
   Prof_FEC.Data[3729] := 47.073;
   Prof_FEC.Data[3730] := 45.575;
   Prof_FEC.Data[3731] := 49.707;
   Prof_FEC.Data[3732] := 41.139;
   Prof_FEC.Data[3733] := 42.988;
   Prof_FEC.Data[3734] := 42.071;
   Prof_FEC.Data[3735] := 46.696;
   Prof_FEC.Data[3736] := 48.281;
   Prof_FEC.Data[3737] := 50.0;
   Prof_FEC.Data[3738] := 47.819;
   Prof_FEC.Data[3739] := 43.092;
   Prof_FEC.Data[3740] := 39.113;
   Prof_FEC.Data[3741] := 42.162;
   Prof_FEC.Data[3742] := 38.882;
   Prof_FEC.Data[3743] := 40.725;
   Prof_FEC.Data[3744] := 45.967;
   Prof_FEC.Data[3745] := 44.621;
   Prof_FEC.Data[3746] := 42.657;
   Prof_FEC.Data[3747] := 41.691;
   Prof_FEC.Data[3748] := 38.553;
   Prof_FEC.Data[3749] := 36.7;
   Prof_FEC.Data[3750] := 41.174;
   Prof_FEC.Data[3751] := 42.239;
   Prof_FEC.Data[3752] := 44.536;
   Prof_FEC.Data[3753] := 45.579;
   Prof_FEC.Data[3754] := 44.151;
   Prof_FEC.Data[3755] := 45.589;
   Prof_FEC.Data[3756] := 37.286;
   Prof_FEC.Data[3757] := 38.42;
   Prof_FEC.Data[3758] := 39.736;
   Prof_FEC.Data[3759] := 40.083;
   Prof_FEC.Data[3760] := 43.392;
   Prof_FEC.Data[3761] := 43.432;
   Prof_FEC.Data[3762] := 44.567;
   Prof_FEC.Data[3763] := 41.102;
   Prof_FEC.Data[3764] := 258.32;
   Prof_FEC.Data[3765] := 265.42;
   Prof_FEC.Data[3766] := 274.62;
   Prof_FEC.Data[3767] := 283.66;
   Prof_FEC.Data[3768] := 322.75;
   Prof_FEC.Data[3769] := 304.51;
   Prof_FEC.Data[3770] := 300.78;
   Prof_FEC.Data[3771] := 303.57;
   Prof_FEC.Data[3772] := 234.61;
   Prof_FEC.Data[3773] := 213.25;
   Prof_FEC.Data[3774] := 207.57;
   Prof_FEC.Data[3775] := 174.41;
   Prof_FEC.Data[3776] := 158.56;
   Prof_FEC.Data[3777] := 195.08;
   Prof_FEC.Data[3778] := 189.59;
   Prof_FEC.Data[3779] := 185.6;
   Prof_FEC.Data[3780] := 140.15;
   Prof_FEC.Data[3781] := 140.92;
   Prof_FEC.Data[3782] := 121.82;
   Prof_FEC.Data[3783] := 137.36;
   Prof_FEC.Data[3784] := 160.3;
   Prof_FEC.Data[3785] := 167.11;
   Prof_FEC.Data[3786] := 179.72;
   Prof_FEC.Data[3787] := 171.92;
   Prof_FEC.Data[3788] := 157.96;
   Prof_FEC.Data[3789] := 131.9;
   Prof_FEC.Data[3790] := 115.89;
   Prof_FEC.Data[3791] := 137.18;
   Prof_FEC.Data[3792] := 197.41;
   Prof_FEC.Data[3793] := 182.04;
   Prof_FEC.Data[3794] := 174.48;
   Prof_FEC.Data[3795] := 154.09;
   Prof_FEC.Data[3796] := 147.21;
   Prof_FEC.Data[3797] := 114.56;
   Prof_FEC.Data[3798] := 135.07;
   Prof_FEC.Data[3799] := 143.52;
   Prof_FEC.Data[3800] := 156.6;
   Prof_FEC.Data[3801] := 175.06;
   Prof_FEC.Data[3802] := 169.73;
   Prof_FEC.Data[3803] := 158.49;
   Prof_FEC.Data[3804] := 155.84;
   Prof_FEC.Data[3805] := 145.64;
   Prof_FEC.Data[3806] := 151.14;
   Prof_FEC.Data[3807] := 155.64;
   Prof_FEC.Data[3808] := 173.23;
   Prof_FEC.Data[3809] := 200.86;
   Prof_FEC.Data[3810] := 202.44;
   Prof_FEC.Data[3811] := 228.82;
   Prof_FEC.Data[3812] := 259.76;
   Prof_FEC.Data[3813] := 299.99;
   Prof_FEC.Data[3814] := 289.9;
   Prof_FEC.Data[3815] := 312.38;
   Prof_FEC.Data[3816] := 349.59;
   Prof_FEC.Data[3817] := 318.2;
   Prof_FEC.Data[3818] := 328.63;
   Prof_FEC.Data[3819] := 318.62;
   Prof_FEC.Data[3820] := 44.911;
   Prof_FEC.Data[3821] := 44.03;
   Prof_FEC.Data[3822] := 43.278;
   Prof_FEC.Data[3823] := 44.686;
   Prof_FEC.Data[3824] := 49.828;
   Prof_FEC.Data[3825] := 50.0;
   Prof_FEC.Data[3826] := 49.932;
   Prof_FEC.Data[3827] := 50.0;
   Prof_FEC.Data[3828] := 47.539;
   Prof_FEC.Data[3829] := 45.295;
   Prof_FEC.Data[3830] := 41.563;
   Prof_FEC.Data[3831] := 45.763;
   Prof_FEC.Data[3832] := 48.697;
   Prof_FEC.Data[3833] := 47.929;
   Prof_FEC.Data[3834] := 47.138;
   Prof_FEC.Data[3835] := 46.2;
   Prof_FEC.Data[3836] := 46.105;
   Prof_FEC.Data[3837] := 47.253;
   Prof_FEC.Data[3838] := 47.456;
   Prof_FEC.Data[3839] := 44.508;
   Prof_FEC.Data[3840] := 46.4;
   Prof_FEC.Data[3841] := 49.261;
   Prof_FEC.Data[3842] := 49.962;
   Prof_FEC.Data[3843] := 45.439;
   Prof_FEC.Data[3844] := 44.952;
   Prof_FEC.Data[3845] := 46.186;
   Prof_FEC.Data[3846] := 41.533;
   Prof_FEC.Data[3847] := 44.847;
   Prof_FEC.Data[3848] := 42.927;
   Prof_FEC.Data[3849] := 45.898;
   Prof_FEC.Data[3850] := 46.995;
   Prof_FEC.Data[3851] := 43.451;
   Prof_FEC.Data[3852] := 41.924;
   Prof_FEC.Data[3853] := 43.779;
   Prof_FEC.Data[3854] := 42.851;
   Prof_FEC.Data[3855] := 42.188;
   Prof_FEC.Data[3856] := 45.768;
   Prof_FEC.Data[3857] := 49.887;
   Prof_FEC.Data[3858] := 47.87;
   Prof_FEC.Data[3859] := 45.856;
   Prof_FEC.Data[3860] := 263.76;
   Prof_FEC.Data[3861] := 229.15;
   Prof_FEC.Data[3862] := 276.0;
   Prof_FEC.Data[3863] := 301.11;
   Prof_FEC.Data[3864] := 346.47;
   Prof_FEC.Data[3865] := 396.8;
   Prof_FEC.Data[3866] := 433.73;
   Prof_FEC.Data[3867] := 448.04;
   Prof_FEC.Data[3868] := 546.36;
   Prof_FEC.Data[3869] := 568.27;
   Prof_FEC.Data[3870] := 566.05;
   Prof_FEC.Data[3871] := 550.87;
   Prof_FEC.Data[3872] := 546.55;
   Prof_FEC.Data[3873] := 682.46;
   Prof_FEC.Data[3874] := 615.99;
   Prof_FEC.Data[3875] := 644.9;
   Prof_FEC.Data[3876] := 616.45;
   Prof_FEC.Data[3877] := 661.92;
   Prof_FEC.Data[3878] := 703.1;
   Prof_FEC.Data[3879] := 715.3;
   Prof_FEC.Data[3880] := 716.63;
   Prof_FEC.Data[3881] := 701.07;
   Prof_FEC.Data[3882] := 690.02;
   Prof_FEC.Data[3883] := 725.13;
   Prof_FEC.Data[3884] := 665.44;
   Prof_FEC.Data[3885] := 718.92;
   Prof_FEC.Data[3886] := 740.98;
   Prof_FEC.Data[3887] := 714.37;
   Prof_FEC.Data[3888] := 714.8;
   Prof_FEC.Data[3889] := 668.72;
   Prof_FEC.Data[3890] := 674.48;
   Prof_FEC.Data[3891] := 631.71;
   Prof_FEC.Data[3892] := 737.7;
   Prof_FEC.Data[3893] := 682.34;
   Prof_FEC.Data[3894] := 714.56;
   Prof_FEC.Data[3895] := 706.64;
   Prof_FEC.Data[3896] := 686.61;
   Prof_FEC.Data[3897] := 642.99;
   Prof_FEC.Data[3898] := 721.74;
   Prof_FEC.Data[3899] := 684.78;
   Prof_FEC.Data[3900] := 734.55;
   Prof_FEC.Data[3901] := 736.82;
   Prof_FEC.Data[3902] := 739.28;
   Prof_FEC.Data[3903] := 650.9;
   Prof_FEC.Data[3904] := 735.17;
   Prof_FEC.Data[3905] := 665.12;
   Prof_FEC.Data[3906] := 713.09;
   Prof_FEC.Data[3907] := 600.1;
   Prof_FEC.Data[3908] := 431.27;
   Prof_FEC.Data[3909] := 355.17;
   Prof_FEC.Data[3910] := 329.2;
   Prof_FEC.Data[3911] := 277.59;
   Prof_FEC.Data[3912] := 255.52;
   Prof_FEC.Data[3913] := 234.2;
   Prof_FEC.Data[3914] := 216.93;
   Prof_FEC.Data[3915] := 236.62;
   Prof_FEC.Data[3916] := 46.915;
   Prof_FEC.Data[3917] := 44.663;
   Prof_FEC.Data[3918] := 45.435;
   Prof_FEC.Data[3919] := 43.41;
   Prof_FEC.Data[3920] := 41.934;
   Prof_FEC.Data[3921] := 41.672;
   Prof_FEC.Data[3922] := 41.871;
   Prof_FEC.Data[3923] := 39.408;
   Prof_FEC.Data[3924] := 45.599;
   Prof_FEC.Data[3925] := 47.848;
   Prof_FEC.Data[3926] := 43.763;
   Prof_FEC.Data[3927] := 44.627;
   Prof_FEC.Data[3928] := 45.059;
   Prof_FEC.Data[3929] := 40.984;
   Prof_FEC.Data[3930] := 43.929;
   Prof_FEC.Data[3931] := 50.0;
   Prof_FEC.Data[3932] := 47.327;
   Prof_FEC.Data[3933] := 47.765;
   Prof_FEC.Data[3934] := 48.227;
   Prof_FEC.Data[3935] := 46.239;
   Prof_FEC.Data[3936] := 43.121;
   Prof_FEC.Data[3937] := 39.625;
   Prof_FEC.Data[3938] := 43.639;
   Prof_FEC.Data[3939] := 44.396;
   Prof_FEC.Data[3940] := 44.924;
   Prof_FEC.Data[3941] := 49.063;
   Prof_FEC.Data[3942] := 49.355;
   Prof_FEC.Data[3943] := 46.777;
   Prof_FEC.Data[3944] := 43.758;
   Prof_FEC.Data[3945] := 40.714;
   Prof_FEC.Data[3946] := 42.239;
   Prof_FEC.Data[3947] := 40.567;
   Prof_FEC.Data[3948] := 43.113;
   Prof_FEC.Data[3949] := 50.0;
   Prof_FEC.Data[3950] := 50.0;
   Prof_FEC.Data[3951] := 44.568;
   Prof_FEC.Data[3952] := 45.219;
   Prof_FEC.Data[3953] := 45.464;
   Prof_FEC.Data[3954] := 45.63;
   Prof_FEC.Data[3955] := 45.472;
   Prof_FEC.Data[3956] := 356.56;
   Prof_FEC.Data[3957] := 321.49;
   Prof_FEC.Data[3958] := 317.85;
   Prof_FEC.Data[3959] := 325.02;
   Prof_FEC.Data[3960] := 387.83;
   Prof_FEC.Data[3961] := 396.37;
   Prof_FEC.Data[3962] := 414.3;
   Prof_FEC.Data[3963] := 445.66;
   Prof_FEC.Data[3964] := 476.39;
   Prof_FEC.Data[3965] := 466.57;
   Prof_FEC.Data[3966] := 556.75;
   Prof_FEC.Data[3967] := 592.06;
   Prof_FEC.Data[3968] := 579.33;
   Prof_FEC.Data[3969] := 630.13;
   Prof_FEC.Data[3970] := 690.21;
   Prof_FEC.Data[3971] := 635.46;
   Prof_FEC.Data[3972] := 664.99;
   Prof_FEC.Data[3973] := 689.12;
   Prof_FEC.Data[3974] := 687.91;
   Prof_FEC.Data[3975] := 703.89;
   Prof_FEC.Data[3976] := 738.22;
   Prof_FEC.Data[3977] := 789.79;
   Prof_FEC.Data[3978] := 750.53;
   Prof_FEC.Data[3979] := 767.52;
   Prof_FEC.Data[3980] := 730.27;
   Prof_FEC.Data[3981] := 715.13;
   Prof_FEC.Data[3982] := 721.37;
   Prof_FEC.Data[3983] := 651.97;
   Prof_FEC.Data[3984] := 759.67;
   Prof_FEC.Data[3985] := 712.24;
   Prof_FEC.Data[3986] := 636.52;
   Prof_FEC.Data[3987] := 718.81;
   Prof_FEC.Data[3988] := 714.57;
   Prof_FEC.Data[3989] := 749.05;
   Prof_FEC.Data[3990] := 676.82;
   Prof_FEC.Data[3991] := 744.38;
   Prof_FEC.Data[3992] := 684.96;
   Prof_FEC.Data[3993] := 726.37;
   Prof_FEC.Data[3994] := 725.06;
   Prof_FEC.Data[3995] := 712.35;
   Prof_FEC.Data[3996] := 686.07;
   Prof_FEC.Data[3997] := 698.41;
   Prof_FEC.Data[3998] := 685.09;
   Prof_FEC.Data[3999] := 685.6;
   Prof_FEC.Data[4000] := 783.53;
   Prof_FEC.Data[4001] := 702.28;
   Prof_FEC.Data[4002] := 695.36;
   Prof_FEC.Data[4003] := 607.19;
   Prof_FEC.Data[4004] := 483.87;
   Prof_FEC.Data[4005] := 365.0;
   Prof_FEC.Data[4006] := 336.72;
   Prof_FEC.Data[4007] := 300.78;
   Prof_FEC.Data[4008] := 286.93;
   Prof_FEC.Data[4009] := 285.94;
   Prof_FEC.Data[4010] := 289.59;
   Prof_FEC.Data[4011] := 269.8;
   Prof_FEC.Data[4012] := 46.807;
   Prof_FEC.Data[4013] := 48.774;
   Prof_FEC.Data[4014] := 50.0;
   Prof_FEC.Data[4015] := 49.332;
   Prof_FEC.Data[4016] := 47.876;
   Prof_FEC.Data[4017] := 46.058;
   Prof_FEC.Data[4018] := 47.326;
   Prof_FEC.Data[4019] := 46.118;
   Prof_FEC.Data[4020] := 50.0;
   Prof_FEC.Data[4021] := 50.0;
   Prof_FEC.Data[4022] := 48.772;
   Prof_FEC.Data[4023] := 48.138;
   Prof_FEC.Data[4024] := 44.613;
   Prof_FEC.Data[4025] := 44.187;
   Prof_FEC.Data[4026] := 47.695;
   Prof_FEC.Data[4027] := 45.371;
   Prof_FEC.Data[4028] := 47.22;
   Prof_FEC.Data[4029] := 48.058;
   Prof_FEC.Data[4030] := 47.997;
   Prof_FEC.Data[4031] := 49.961;
   Prof_FEC.Data[4032] := 48.472;
   Prof_FEC.Data[4033] := 46.735;
   Prof_FEC.Data[4034] := 48.774;
   Prof_FEC.Data[4035] := 48.154;
   Prof_FEC.Data[4036] := 49.892;
   Prof_FEC.Data[4037] := 50.0;
   Prof_FEC.Data[4038] := 50.0;
   Prof_FEC.Data[4039] := 50.0;
   Prof_FEC.Data[4040] := 48.64;
   Prof_FEC.Data[4041] := 49.155;
   Prof_FEC.Data[4042] := 48.249;
   Prof_FEC.Data[4043] := 50.0;
   Prof_FEC.Data[4044] := 50.0;
   Prof_FEC.Data[4045] := 50.0;
   Prof_FEC.Data[4046] := 50.0;
   Prof_FEC.Data[4047] := 50.0;
   Prof_FEC.Data[4048] := 49.777;
   Prof_FEC.Data[4049] := 49.517;
   Prof_FEC.Data[4050] := 45.302;
   Prof_FEC.Data[4051] := 46.794;
   Prof_FEC.Data[4052] := 298.02;
   Prof_FEC.Data[4053] := 348.75;
   Prof_FEC.Data[4054] := 351.67;
   Prof_FEC.Data[4055] := 385.15;
   Prof_FEC.Data[4056] := 352.57;
   Prof_FEC.Data[4057] := 355.72;
   Prof_FEC.Data[4058] := 331.72;
   Prof_FEC.Data[4059] := 426.49;
   Prof_FEC.Data[4060] := 423.58;
   Prof_FEC.Data[4061] := 484.85;
   Prof_FEC.Data[4062] := 478.55;
   Prof_FEC.Data[4063] := 444.25;
   Prof_FEC.Data[4064] := 463.66;
   Prof_FEC.Data[4065] := 542.66;
   Prof_FEC.Data[4066] := 577.83;
   Prof_FEC.Data[4067] := 510.24;
   Prof_FEC.Data[4068] := 585.58;
   Prof_FEC.Data[4069] := 583.65;
   Prof_FEC.Data[4070] := 567.73;
   Prof_FEC.Data[4071] := 596.88;
   Prof_FEC.Data[4072] := 671.0;
   Prof_FEC.Data[4073] := 670.74;
   Prof_FEC.Data[4074] := 640.55;
   Prof_FEC.Data[4075] := 703.92;
   Prof_FEC.Data[4076] := 651.03;
   Prof_FEC.Data[4077] := 604.1;
   Prof_FEC.Data[4078] := 648.04;
   Prof_FEC.Data[4079] := 619.02;
   Prof_FEC.Data[4080] := 590.62;
   Prof_FEC.Data[4081] := 569.72;
   Prof_FEC.Data[4082] := 564.26;
   Prof_FEC.Data[4083] := 548.4;
   Prof_FEC.Data[4084] := 607.0;
   Prof_FEC.Data[4085] := 630.15;
   Prof_FEC.Data[4086] := 573.76;
   Prof_FEC.Data[4087] := 544.51;
   Prof_FEC.Data[4088] := 531.38;
   Prof_FEC.Data[4089] := 601.3;
   Prof_FEC.Data[4090] := 552.9;
   Prof_FEC.Data[4091] := 677.9;
   Prof_FEC.Data[4092] := 693.65;
   Prof_FEC.Data[4093] := 593.99;
   Prof_FEC.Data[4094] := 560.46;
   Prof_FEC.Data[4095] := 653.74;
   Prof_FEC.Data[4096] := 740.86;
   Prof_FEC.Data[4097] := 626.23;
   Prof_FEC.Data[4098] := 682.94;
   Prof_FEC.Data[4099] := 481.66;
   Prof_FEC.Data[4100] := 393.42;
   Prof_FEC.Data[4101] := 373.99;
   Prof_FEC.Data[4102] := 346.88;
   Prof_FEC.Data[4103] := 309.67;
   Prof_FEC.Data[4104] := 296.54;
   Prof_FEC.Data[4105] := 288.07;
   Prof_FEC.Data[4106] := 289.18;
   Prof_FEC.Data[4107] := 280.45;
   Prof_FEC.Data[4108] := 46.042;
   Prof_FEC.Data[4109] := 50.0;
   Prof_FEC.Data[4110] := 50.0;
   Prof_FEC.Data[4111] := 49.808;
   Prof_FEC.Data[4112] := 45.426;
   Prof_FEC.Data[4113] := 46.312;
   Prof_FEC.Data[4114] := 43.196;
   Prof_FEC.Data[4115] := 46.23;
   Prof_FEC.Data[4116] := 50.0;
   Prof_FEC.Data[4117] := 50.0;
   Prof_FEC.Data[4118] := 50.0;
   Prof_FEC.Data[4119] := 47.566;
   Prof_FEC.Data[4120] := 46.692;
   Prof_FEC.Data[4121] := 46.043;
   Prof_FEC.Data[4122] := 44.113;
   Prof_FEC.Data[4123] := 43.549;
   Prof_FEC.Data[4124] := 48.932;
   Prof_FEC.Data[4125] := 46.072;
   Prof_FEC.Data[4126] := 44.029;
   Prof_FEC.Data[4127] := 42.86;
   Prof_FEC.Data[4128] := 46.235;
   Prof_FEC.Data[4129] := 44.883;
   Prof_FEC.Data[4130] := 43.177;
   Prof_FEC.Data[4131] := 43.567;
   Prof_FEC.Data[4132] := 46.452;
   Prof_FEC.Data[4133] := 46.155;
   Prof_FEC.Data[4134] := 47.375;
   Prof_FEC.Data[4135] := 45.482;
   Prof_FEC.Data[4136] := 43.393;
   Prof_FEC.Data[4137] := 40.504;
   Prof_FEC.Data[4138] := 45.073;
   Prof_FEC.Data[4139] := 45.076;
   Prof_FEC.Data[4140] := 43.295;
   Prof_FEC.Data[4141] := 45.415;
   Prof_FEC.Data[4142] := 42.79;
   Prof_FEC.Data[4143] := 42.803;
   Prof_FEC.Data[4144] := 37.454;
   Prof_FEC.Data[4145] := 40.137;
   Prof_FEC.Data[4146] := 40.222;
   Prof_FEC.Data[4147] := 43.649;
   Prof_FEC.Data[4148] := 298.38;
   Prof_FEC.Data[4149] := 317.4;
   Prof_FEC.Data[4150] := 335.28;
   Prof_FEC.Data[4151] := 348.28;
   Prof_FEC.Data[4152] := 404.41;
   Prof_FEC.Data[4153] := 439.44;
   Prof_FEC.Data[4154] := 422.26;
   Prof_FEC.Data[4155] := 470.06;
   Prof_FEC.Data[4156] := 475.74;
   Prof_FEC.Data[4157] := 502.16;
   Prof_FEC.Data[4158] := 466.84;
   Prof_FEC.Data[4159] := 542.1;
   Prof_FEC.Data[4160] := 572.83;
   Prof_FEC.Data[4161] := 578.28;
   Prof_FEC.Data[4162] := 584.98;
   Prof_FEC.Data[4163] := 542.46;
   Prof_FEC.Data[4164] := 574.9;
   Prof_FEC.Data[4165] := 609.15;
   Prof_FEC.Data[4166] := 590.4;
   Prof_FEC.Data[4167] := 623.75;
   Prof_FEC.Data[4168] := 712.72;
   Prof_FEC.Data[4169] := 595.76;
   Prof_FEC.Data[4170] := 620.48;
   Prof_FEC.Data[4171] := 690.37;
   Prof_FEC.Data[4172] := 668.89;
   Prof_FEC.Data[4173] := 669.89;
   Prof_FEC.Data[4174] := 645.78;
   Prof_FEC.Data[4175] := 694.32;
   Prof_FEC.Data[4176] := 568.53;
   Prof_FEC.Data[4177] := 626.3;
   Prof_FEC.Data[4178] := 603.87;
   Prof_FEC.Data[4179] := 579.81;
   Prof_FEC.Data[4180] := 617.55;
   Prof_FEC.Data[4181] := 624.83;
   Prof_FEC.Data[4182] := 641.48;
   Prof_FEC.Data[4183] := 687.35;
   Prof_FEC.Data[4184] := 604.7;
   Prof_FEC.Data[4185] := 622.94;
   Prof_FEC.Data[4186] := 621.68;
   Prof_FEC.Data[4187] := 608.58;
   Prof_FEC.Data[4188] := 677.04;
   Prof_FEC.Data[4189] := 596.59;
   Prof_FEC.Data[4190] := 536.13;
   Prof_FEC.Data[4191] := 610.02;
   Prof_FEC.Data[4192] := 607.73;
   Prof_FEC.Data[4193] := 628.47;
   Prof_FEC.Data[4194] := 604.46;
   Prof_FEC.Data[4195] := 556.36;
   Prof_FEC.Data[4196] := 422.99;
   Prof_FEC.Data[4197] := 331.35;
   Prof_FEC.Data[4198] := 301.77;
   Prof_FEC.Data[4199] := 247.68;
   Prof_FEC.Data[4200] := 251.56;
   Prof_FEC.Data[4201] := 230.63;
   Prof_FEC.Data[4202] := 251.45;
   Prof_FEC.Data[4203] := 249.56;
   Prof_FEC.Data[4204] := 42.584;
   Prof_FEC.Data[4205] := 45.646;
   Prof_FEC.Data[4206] := 45.154;
   Prof_FEC.Data[4207] := 40.895;
   Prof_FEC.Data[4208] := 43.575;
   Prof_FEC.Data[4209] := 42.58;
   Prof_FEC.Data[4210] := 41.636;
   Prof_FEC.Data[4211] := 43.009;
   Prof_FEC.Data[4212] := 43.941;
   Prof_FEC.Data[4213] := 41.672;
   Prof_FEC.Data[4214] := 45.951;
   Prof_FEC.Data[4215] := 45.261;
   Prof_FEC.Data[4216] := 43.426;
   Prof_FEC.Data[4217] := 40.64;
   Prof_FEC.Data[4218] := 43.438;
   Prof_FEC.Data[4219] := 41.021;
   Prof_FEC.Data[4220] := 44.548;
   Prof_FEC.Data[4221] := 46.217;
   Prof_FEC.Data[4222] := 43.932;
   Prof_FEC.Data[4223] := 45.155;
   Prof_FEC.Data[4224] := 41.42;
   Prof_FEC.Data[4225] := 40.693;
   Prof_FEC.Data[4226] := 39.776;
   Prof_FEC.Data[4227] := 43.119;
   Prof_FEC.Data[4228] := 46.806;
   Prof_FEC.Data[4229] := 42.925;
   Prof_FEC.Data[4230] := 43.398;
   Prof_FEC.Data[4231] := 45.375;
   Prof_FEC.Data[4232] := 41.858;
   Prof_FEC.Data[4233] := 41.765;
   Prof_FEC.Data[4234] := 42.076;
   Prof_FEC.Data[4235] := 39.465;
   Prof_FEC.Data[4236] := 43.627;
   Prof_FEC.Data[4237] := 41.576;
   Prof_FEC.Data[4238] := 43.878;
   Prof_FEC.Data[4239] := 39.875;
   Prof_FEC.Data[4240] := 41.185;
   Prof_FEC.Data[4241] := 38.026;
   Prof_FEC.Data[4242] := 40.587;
   Prof_FEC.Data[4243] := 38.997;
   Prof_FEC.Data[4244] := 228.78;
   Prof_FEC.Data[4245] := 262.94;
   Prof_FEC.Data[4246] := 237.14;
   Prof_FEC.Data[4247] := 296.3;
   Prof_FEC.Data[4248] := 336.89;
   Prof_FEC.Data[4249] := 353.55;
   Prof_FEC.Data[4250] := 378.06;
   Prof_FEC.Data[4251] := 417.63;
   Prof_FEC.Data[4252] := 450.82;
   Prof_FEC.Data[4253] := 462.32;
   Prof_FEC.Data[4254] := 503.17;
   Prof_FEC.Data[4255] := 498.35;
   Prof_FEC.Data[4256] := 529.09;
   Prof_FEC.Data[4257] := 548.23;
   Prof_FEC.Data[4258] := 508.56;
   Prof_FEC.Data[4259] := 582.94;
   Prof_FEC.Data[4260] := 552.39;
   Prof_FEC.Data[4261] := 542.81;
   Prof_FEC.Data[4262] := 565.52;
   Prof_FEC.Data[4263] := 565.86;
   Prof_FEC.Data[4264] := 589.08;
   Prof_FEC.Data[4265] := 602.75;
   Prof_FEC.Data[4266] := 626.59;
   Prof_FEC.Data[4267] := 683.92;
   Prof_FEC.Data[4268] := 690.51;
   Prof_FEC.Data[4269] := 653.86;
   Prof_FEC.Data[4270] := 655.36;
   Prof_FEC.Data[4271] := 597.4;
   Prof_FEC.Data[4272] := 525.74;
   Prof_FEC.Data[4273] := 517.07;
   Prof_FEC.Data[4274] := 527.9;
   Prof_FEC.Data[4275] := 546.92;
   Prof_FEC.Data[4276] := 501.56;
   Prof_FEC.Data[4277] := 545.48;
   Prof_FEC.Data[4278] := 596.96;
   Prof_FEC.Data[4279] := 483.72;
   Prof_FEC.Data[4280] := 562.08;
   Prof_FEC.Data[4281] := 488.63;
   Prof_FEC.Data[4282] := 599.12;
   Prof_FEC.Data[4283] := 553.38;
   Prof_FEC.Data[4284] := 568.25;
   Prof_FEC.Data[4285] := 595.77;
   Prof_FEC.Data[4286] := 543.28;
   Prof_FEC.Data[4287] := 621.11;
   Prof_FEC.Data[4288] := 555.95;
   Prof_FEC.Data[4289] := 623.5;
   Prof_FEC.Data[4290] := 530.62;
   Prof_FEC.Data[4291] := 468.19;
   Prof_FEC.Data[4292] := 338.82;
   Prof_FEC.Data[4293] := 267.64;
   Prof_FEC.Data[4294] := 258.63;
   Prof_FEC.Data[4295] := 252.06;
   Prof_FEC.Data[4296] := 271.73;
   Prof_FEC.Data[4297] := 219.33;
   Prof_FEC.Data[4298] := 203.92;
   Prof_FEC.Data[4299] := 216.48;
   Prof_FEC.Data[4300] := 40.964;
   Prof_FEC.Data[4301] := 39.859;
   Prof_FEC.Data[4302] := 38.9;
   Prof_FEC.Data[4303] := 38.015;
   Prof_FEC.Data[4304] := 38.925;
   Prof_FEC.Data[4305] := 39.321;
   Prof_FEC.Data[4306] := 37.614;
   Prof_FEC.Data[4307] := 38.837;
   Prof_FEC.Data[4308] := 40.842;
   Prof_FEC.Data[4309] := 39.534;
   Prof_FEC.Data[4310] := 43.164;
   Prof_FEC.Data[4311] := 42.305;
   Prof_FEC.Data[4312] := 38.735;
   Prof_FEC.Data[4313] := 39.378;
   Prof_FEC.Data[4314] := 38.896;
   Prof_FEC.Data[4315] := 38.237;
   Prof_FEC.Data[4316] := 41.62;
   Prof_FEC.Data[4317] := 42.827;
   Prof_FEC.Data[4318] := 40.415;
   Prof_FEC.Data[4319] := 42.696;
   Prof_FEC.Data[4320] := 40.915;
   Prof_FEC.Data[4321] := 42.188;
   Prof_FEC.Data[4322] := 42.927;
   Prof_FEC.Data[4323] := 43.594;
   Prof_FEC.Data[4324] := 44.611;
   Prof_FEC.Data[4325] := 46.489;
   Prof_FEC.Data[4326] := 48.803;
   Prof_FEC.Data[4327] := 42.237;
   Prof_FEC.Data[4328] := 44.559;
   Prof_FEC.Data[4329] := 42.739;
   Prof_FEC.Data[4330] := 43.823;
   Prof_FEC.Data[4331] := 43.105;
   Prof_FEC.Data[4332] := 44.611;
   Prof_FEC.Data[4333] := 46.543;
   Prof_FEC.Data[4334] := 44.644;
   Prof_FEC.Data[4335] := 43.431;
   Prof_FEC.Data[4336] := 45.935;
   Prof_FEC.Data[4337] := 44.609;
   Prof_FEC.Data[4338] := 42.329;
   Prof_FEC.Data[4339] := 42.1;
   Prof_FEC.Data[4340] := 298.58;
   Prof_FEC.Data[4341] := 313.24;
   Prof_FEC.Data[4342] := 312.75;
   Prof_FEC.Data[4343] := 284.72;
   Prof_FEC.Data[4344] := 280.98;
   Prof_FEC.Data[4345] := 294.6;
   Prof_FEC.Data[4346] := 278.06;
   Prof_FEC.Data[4347] := 296.58;
   Prof_FEC.Data[4348] := 286.73;
   Prof_FEC.Data[4349] := 299.13;
   Prof_FEC.Data[4350] := 325.73;
   Prof_FEC.Data[4351] := 311.08;
   Prof_FEC.Data[4352] := 262.82;
   Prof_FEC.Data[4353] := 245.95;
   Prof_FEC.Data[4354] := 242.28;
   Prof_FEC.Data[4355] := 270.88;
   Prof_FEC.Data[4356] := 268.75;
   Prof_FEC.Data[4357] := 356.64;
   Prof_FEC.Data[4358] := 351.15;
   Prof_FEC.Data[4359] := 360.61;
   Prof_FEC.Data[4360] := 349.96;
   Prof_FEC.Data[4361] := 325.1;
   Prof_FEC.Data[4362] := 340.06;
   Prof_FEC.Data[4363] := 397.32;
   Prof_FEC.Data[4364] := 371.79;
   Prof_FEC.Data[4365] := 395.48;
   Prof_FEC.Data[4366] := 345.22;
   Prof_FEC.Data[4367] := 328.57;
   Prof_FEC.Data[4368] := 275.55;
   Prof_FEC.Data[4369] := 255.33;
   Prof_FEC.Data[4370] := 237.66;
   Prof_FEC.Data[4371] := 268.04;
   Prof_FEC.Data[4372] := 297.33;
   Prof_FEC.Data[4373] := 266.42;
   Prof_FEC.Data[4374] := 261.27;
   Prof_FEC.Data[4375] := 240.4;
   Prof_FEC.Data[4376] := 238.57;
   Prof_FEC.Data[4377] := 274.52;
   Prof_FEC.Data[4378] := 240.93;
   Prof_FEC.Data[4379] := 251.06;
   Prof_FEC.Data[4380] := 289.05;
   Prof_FEC.Data[4381] := 246.35;
   Prof_FEC.Data[4382] := 244.95;
   Prof_FEC.Data[4383] := 201.86;
   Prof_FEC.Data[4384] := 139.79;
   Prof_FEC.Data[4385] := 123.58;
   Prof_FEC.Data[4386] := 122.73;
   Prof_FEC.Data[4387] := 137.01;
   Prof_FEC.Data[4388] := 193.76;
   Prof_FEC.Data[4389] := 213.89;
   Prof_FEC.Data[4390] := 222.18;
   Prof_FEC.Data[4391] := 256.95;
   Prof_FEC.Data[4392] := 278.46;
   Prof_FEC.Data[4393] := 262.26;
   Prof_FEC.Data[4394] := 318.89;
   Prof_FEC.Data[4395] := 306.67;
   Prof_FEC.Data[4396] := 44.037;
   Prof_FEC.Data[4397] := 45.845;
   Prof_FEC.Data[4398] := 42.133;
   Prof_FEC.Data[4399] := 43.183;
   Prof_FEC.Data[4400] := 47.919;
   Prof_FEC.Data[4401] := 46.074;
   Prof_FEC.Data[4402] := 48.49;
   Prof_FEC.Data[4403] := 49.003;
   Prof_FEC.Data[4404] := 46.148;
   Prof_FEC.Data[4405] := 45.146;
   Prof_FEC.Data[4406] := 43.483;
   Prof_FEC.Data[4407] := 42.543;
   Prof_FEC.Data[4408] := 43.633;
   Prof_FEC.Data[4409] := 44.526;
   Prof_FEC.Data[4410] := 41.504;
   Prof_FEC.Data[4411] := 46.006;
   Prof_FEC.Data[4412] := 41.017;
   Prof_FEC.Data[4413] := 42.429;
   Prof_FEC.Data[4414] := 40.954;
   Prof_FEC.Data[4415] := 39.75;
   Prof_FEC.Data[4416] := 45.931;
   Prof_FEC.Data[4417] := 47.108;
   Prof_FEC.Data[4418] := 42.567;
   Prof_FEC.Data[4419] := 44.458;
   Prof_FEC.Data[4420] := 44.842;
   Prof_FEC.Data[4421] := 41.047;
   Prof_FEC.Data[4422] := 40.391;
   Prof_FEC.Data[4423] := 42.682;
   Prof_FEC.Data[4424] := 44.165;
   Prof_FEC.Data[4425] := 45.166;
   Prof_FEC.Data[4426] := 44.773;
   Prof_FEC.Data[4427] := 44.563;
   Prof_FEC.Data[4428] := 40.737;
   Prof_FEC.Data[4429] := 42.922;
   Prof_FEC.Data[4430] := 41.722;
   Prof_FEC.Data[4431] := 42.969;
   Prof_FEC.Data[4432] := 41.411;
   Prof_FEC.Data[4433] := 44.003;
   Prof_FEC.Data[4434] := 46.293;
   Prof_FEC.Data[4435] := 46.085;
   Prof_FEC.Data[4436] := 275.76;
   Prof_FEC.Data[4437] := 266.93;
   Prof_FEC.Data[4438] := 275.02;
   Prof_FEC.Data[4439] := 288.08;
   Prof_FEC.Data[4440] := 371.54;
   Prof_FEC.Data[4441] := 357.21;
   Prof_FEC.Data[4442] := 346.65;
   Prof_FEC.Data[4443] := 293.68;
   Prof_FEC.Data[4444] := 236.87;
   Prof_FEC.Data[4445] := 227.72;
   Prof_FEC.Data[4446] := 219.96;
   Prof_FEC.Data[4447] := 199.09;
   Prof_FEC.Data[4448] := 212.18;
   Prof_FEC.Data[4449] := 205.09;
   Prof_FEC.Data[4450] := 183.07;
   Prof_FEC.Data[4451] := 193.95;
   Prof_FEC.Data[4452] := 167.03;
   Prof_FEC.Data[4453] := 152.5;
   Prof_FEC.Data[4454] := 147.78;
   Prof_FEC.Data[4455] := 143.1;
   Prof_FEC.Data[4456] := 170.36;
   Prof_FEC.Data[4457] := 170.19;
   Prof_FEC.Data[4458] := 175.26;
   Prof_FEC.Data[4459] := 160.24;
   Prof_FEC.Data[4460] := 140.31;
   Prof_FEC.Data[4461] := 114.83;
   Prof_FEC.Data[4462] := 109.81;
   Prof_FEC.Data[4463] := 119.07;
   Prof_FEC.Data[4464] := 148.57;
   Prof_FEC.Data[4465] := 130.36;
   Prof_FEC.Data[4466] := 160.66;
   Prof_FEC.Data[4467] := 143.82;
   Prof_FEC.Data[4468] := 125.45;
   Prof_FEC.Data[4469] := 124.47;
   Prof_FEC.Data[4470] := 117.63;
   Prof_FEC.Data[4471] := 111.37;
   Prof_FEC.Data[4472] := 117.4;
   Prof_FEC.Data[4473] := 145.99;
   Prof_FEC.Data[4474] := 147.28;
   Prof_FEC.Data[4475] := 143.28;
   Prof_FEC.Data[4476] := 132.74;
   Prof_FEC.Data[4477] := 118.04;
   Prof_FEC.Data[4478] := 110.68;
   Prof_FEC.Data[4479] := 123.0;
   Prof_FEC.Data[4480] := 137.57;
   Prof_FEC.Data[4481] := 140.29;
   Prof_FEC.Data[4482] := 142.78;
   Prof_FEC.Data[4483] := 151.53;
   Prof_FEC.Data[4484] := 180.29;
   Prof_FEC.Data[4485] := 207.22;
   Prof_FEC.Data[4486] := 233.52;
   Prof_FEC.Data[4487] := 240.12;
   Prof_FEC.Data[4488] := 266.97;
   Prof_FEC.Data[4489] := 315.69;
   Prof_FEC.Data[4490] := 278.14;
   Prof_FEC.Data[4491] := 316.66;
   Prof_FEC.Data[4492] := 43.143;
   Prof_FEC.Data[4493] := 44.231;
   Prof_FEC.Data[4494] := 43.702;
   Prof_FEC.Data[4495] := 45.205;
   Prof_FEC.Data[4496] := 45.388;
   Prof_FEC.Data[4497] := 46.62;
   Prof_FEC.Data[4498] := 46.595;
   Prof_FEC.Data[4499] := 45.92;
   Prof_FEC.Data[4500] := 44.548;
   Prof_FEC.Data[4501] := 41.69;
   Prof_FEC.Data[4502] := 43.686;
   Prof_FEC.Data[4503] := 42.509;
   Prof_FEC.Data[4504] := 44.076;
   Prof_FEC.Data[4505] := 46.976;
   Prof_FEC.Data[4506] := 47.886;
   Prof_FEC.Data[4507] := 44.741;
   Prof_FEC.Data[4508] := 46.359;
   Prof_FEC.Data[4509] := 41.495;
   Prof_FEC.Data[4510] := 45.405;
   Prof_FEC.Data[4511] := 44.745;
   Prof_FEC.Data[4512] := 46.343;
   Prof_FEC.Data[4513] := 47.895;
   Prof_FEC.Data[4514] := 45.906;
   Prof_FEC.Data[4515] := 47.333;
   Prof_FEC.Data[4516] := 43.493;
   Prof_FEC.Data[4517] := 42.238;
   Prof_FEC.Data[4518] := 40.51;
   Prof_FEC.Data[4519] := 44.783;
   Prof_FEC.Data[4520] := 47.844;
   Prof_FEC.Data[4521] := 46.419;
   Prof_FEC.Data[4522] := 47.08;
   Prof_FEC.Data[4523] := 46.13;
   Prof_FEC.Data[4524] := 43.294;
   Prof_FEC.Data[4525] := 47.501;
   Prof_FEC.Data[4526] := 45.413;
   Prof_FEC.Data[4527] := 43.431;
   Prof_FEC.Data[4528] := 50.0;
   Prof_FEC.Data[4529] := 48.969;
   Prof_FEC.Data[4530] := 47.894;
   Prof_FEC.Data[4531] := 48.406;
   Prof_FEC.Data[4532] := 284.36;
   Prof_FEC.Data[4533] := 276.07;
   Prof_FEC.Data[4534] := 274.73;
   Prof_FEC.Data[4535] := 343.81;
   Prof_FEC.Data[4536] := 399.23;
   Prof_FEC.Data[4537] := 399.58;
   Prof_FEC.Data[4538] := 434.63;
   Prof_FEC.Data[4539] := 431.41;
   Prof_FEC.Data[4540] := 440.86;
   Prof_FEC.Data[4541] := 482.39;
   Prof_FEC.Data[4542] := 562.75;
   Prof_FEC.Data[4543] := 567.19;
   Prof_FEC.Data[4544] := 550.25;
   Prof_FEC.Data[4545] := 584.41;
   Prof_FEC.Data[4546] := 617.29;
   Prof_FEC.Data[4547] := 594.84;
   Prof_FEC.Data[4548] := 601.06;
   Prof_FEC.Data[4549] := 626.98;
   Prof_FEC.Data[4550] := 591.85;
   Prof_FEC.Data[4551] := 615.5;
   Prof_FEC.Data[4552] := 582.5;
   Prof_FEC.Data[4553] := 602.91;
   Prof_FEC.Data[4554] := 662.79;
   Prof_FEC.Data[4555] := 711.39;
   Prof_FEC.Data[4556] := 675.88;
   Prof_FEC.Data[4557] := 644.44;
   Prof_FEC.Data[4558] := 620.67;
   Prof_FEC.Data[4559] := 639.28;
   Prof_FEC.Data[4560] := 598.32;
   Prof_FEC.Data[4561] := 589.98;
   Prof_FEC.Data[4562] := 553.96;
   Prof_FEC.Data[4563] := 501.95;
   Prof_FEC.Data[4564] := 614.72;
   Prof_FEC.Data[4565] := 589.54;
   Prof_FEC.Data[4566] := 610.6;
   Prof_FEC.Data[4567] := 627.34;
   Prof_FEC.Data[4568] := 665.6;
   Prof_FEC.Data[4569] := 649.93;
   Prof_FEC.Data[4570] := 625.73;
   Prof_FEC.Data[4571] := 645.72;
   Prof_FEC.Data[4572] := 712.88;
   Prof_FEC.Data[4573] := 610.77;
   Prof_FEC.Data[4574] := 709.29;
   Prof_FEC.Data[4575] := 683.81;
   Prof_FEC.Data[4576] := 820.42;
   Prof_FEC.Data[4577] := 773.03;
   Prof_FEC.Data[4578] := 727.18;
   Prof_FEC.Data[4579] := 631.87;
   Prof_FEC.Data[4580] := 445.21;
   Prof_FEC.Data[4581] := 341.42;
   Prof_FEC.Data[4582] := 267.52;
   Prof_FEC.Data[4583] := 259.53;
   Prof_FEC.Data[4584] := 247.71;
   Prof_FEC.Data[4585] := 223.27;
   Prof_FEC.Data[4586] := 201.36;
   Prof_FEC.Data[4587] := 262.35;
   Prof_FEC.Data[4588] := 46.445;
   Prof_FEC.Data[4589] := 43.606;
   Prof_FEC.Data[4590] := 45.858;
   Prof_FEC.Data[4591] := 44.226;
   Prof_FEC.Data[4592] := 42.695;
   Prof_FEC.Data[4593] := 42.017;
   Prof_FEC.Data[4594] := 42.569;
   Prof_FEC.Data[4595] := 42.322;
   Prof_FEC.Data[4596] := 46.346;
   Prof_FEC.Data[4597] := 45.202;
   Prof_FEC.Data[4598] := 44.215;
   Prof_FEC.Data[4599] := 46.161;
   Prof_FEC.Data[4600] := 44.135;
   Prof_FEC.Data[4601] := 44.126;
   Prof_FEC.Data[4602] := 45.628;
   Prof_FEC.Data[4603] := 44.056;
   Prof_FEC.Data[4604] := 50.0;
   Prof_FEC.Data[4605] := 50.0;
   Prof_FEC.Data[4606] := 50.0;
   Prof_FEC.Data[4607] := 50.0;
   Prof_FEC.Data[4608] := 47.743;
   Prof_FEC.Data[4609] := 46.52;
   Prof_FEC.Data[4610] := 48.729;
   Prof_FEC.Data[4611] := 48.074;
   Prof_FEC.Data[4612] := 50.0;
   Prof_FEC.Data[4613] := 49.109;
   Prof_FEC.Data[4614] := 50.0;
   Prof_FEC.Data[4615] := 50.0;
   Prof_FEC.Data[4616] := 46.864;
   Prof_FEC.Data[4617] := 45.994;
   Prof_FEC.Data[4618] := 48.063;
   Prof_FEC.Data[4619] := 50.0;
   Prof_FEC.Data[4620] := 49.94;
   Prof_FEC.Data[4621] := 50.0;
   Prof_FEC.Data[4622] := 48.303;
   Prof_FEC.Data[4623] := 49.716;
   Prof_FEC.Data[4624] := 48.983;
   Prof_FEC.Data[4625] := 44.811;
   Prof_FEC.Data[4626] := 43.048;
   Prof_FEC.Data[4627] := 43.571;
   Prof_FEC.Data[4628] := 292.13;
   Prof_FEC.Data[4629] := 317.43;
   Prof_FEC.Data[4630] := 329.52;
   Prof_FEC.Data[4631] := 362.96;
   Prof_FEC.Data[4632] := 386.49;
   Prof_FEC.Data[4633] := 417.31;
   Prof_FEC.Data[4634] := 430.63;
   Prof_FEC.Data[4635] := 466.91;
   Prof_FEC.Data[4636] := 508.25;
   Prof_FEC.Data[4637] := 440.88;
   Prof_FEC.Data[4638] := 447.2;
   Prof_FEC.Data[4639] := 483.75;
   Prof_FEC.Data[4640] := 536.53;
   Prof_FEC.Data[4641] := 558.72;
   Prof_FEC.Data[4642] := 627.09;
   Prof_FEC.Data[4643] := 607.89;
   Prof_FEC.Data[4644] := 676.51;
   Prof_FEC.Data[4645] := 690.37;
   Prof_FEC.Data[4646] := 646.17;
   Prof_FEC.Data[4647] := 744.26;
   Prof_FEC.Data[4648] := 683.63;
   Prof_FEC.Data[4649] := 662.57;
   Prof_FEC.Data[4650] := 664.28;
   Prof_FEC.Data[4651] := 614.81;
   Prof_FEC.Data[4652] := 706.12;
   Prof_FEC.Data[4653] := 665.95;
   Prof_FEC.Data[4654] := 646.47;
   Prof_FEC.Data[4655] := 655.15;
   Prof_FEC.Data[4656] := 619.76;
   Prof_FEC.Data[4657] := 619.63;
   Prof_FEC.Data[4658] := 627.72;
   Prof_FEC.Data[4659] := 554.3;
   Prof_FEC.Data[4660] := 650.8;
   Prof_FEC.Data[4661] := 687.67;
   Prof_FEC.Data[4662] := 653.09;
   Prof_FEC.Data[4663] := 613.3;
   Prof_FEC.Data[4664] := 696.62;
   Prof_FEC.Data[4665] := 669.57;
   Prof_FEC.Data[4666] := 621.81;
   Prof_FEC.Data[4667] := 665.62;
   Prof_FEC.Data[4668] := 653.84;
   Prof_FEC.Data[4669] := 634.95;
   Prof_FEC.Data[4670] := 627.62;
   Prof_FEC.Data[4671] := 697.19;
   Prof_FEC.Data[4672] := 638.92;
   Prof_FEC.Data[4673] := 667.48;
   Prof_FEC.Data[4674] := 703.21;
   Prof_FEC.Data[4675] := 512.79;
   Prof_FEC.Data[4676] := 407.24;
   Prof_FEC.Data[4677] := 311.62;
   Prof_FEC.Data[4678] := 290.42;
   Prof_FEC.Data[4679] := 292.63;
   Prof_FEC.Data[4680] := 262.95;
   Prof_FEC.Data[4681] := 249.05;
   Prof_FEC.Data[4682] := 266.84;
   Prof_FEC.Data[4683] := 251.14;
   Prof_FEC.Data[4684] := 46.954;
   Prof_FEC.Data[4685] := 47.075;
   Prof_FEC.Data[4686] := 44.466;
   Prof_FEC.Data[4687] := 43.58;
   Prof_FEC.Data[4688] := 44.69;
   Prof_FEC.Data[4689] := 41.222;
   Prof_FEC.Data[4690] := 41.45;
   Prof_FEC.Data[4691] := 46.183;
   Prof_FEC.Data[4692] := 45.113;
   Prof_FEC.Data[4693] := 45.539;
   Prof_FEC.Data[4694] := 46.225;
   Prof_FEC.Data[4695] := 44.47;
   Prof_FEC.Data[4696] := 41.361;
   Prof_FEC.Data[4697] := 43.2;
   Prof_FEC.Data[4698] := 44.072;
   Prof_FEC.Data[4699] := 42.92;
   Prof_FEC.Data[4700] := 44.893;
   Prof_FEC.Data[4701] := 48.826;
   Prof_FEC.Data[4702] := 46.842;
   Prof_FEC.Data[4703] := 47.715;
   Prof_FEC.Data[4704] := 46.435;
   Prof_FEC.Data[4705] := 44.782;
   Prof_FEC.Data[4706] := 45.594;
   Prof_FEC.Data[4707] := 45.005;
   Prof_FEC.Data[4708] := 43.413;
   Prof_FEC.Data[4709] := 44.963;
   Prof_FEC.Data[4710] := 46.237;
   Prof_FEC.Data[4711] := 47.435;
   Prof_FEC.Data[4712] := 44.783;
   Prof_FEC.Data[4713] := 41.37;
   Prof_FEC.Data[4714] := 45.497;
   Prof_FEC.Data[4715] := 45.828;
   Prof_FEC.Data[4716] := 48.134;
   Prof_FEC.Data[4717] := 50.0;
   Prof_FEC.Data[4718] := 49.058;
   Prof_FEC.Data[4719] := 47.956;
   Prof_FEC.Data[4720] := 45.708;
   Prof_FEC.Data[4721] := 45.934;
   Prof_FEC.Data[4722] := 45.528;
   Prof_FEC.Data[4723] := 45.239;
   Prof_FEC.Data[4724] := 292.14;
   Prof_FEC.Data[4725] := 287.0;
   Prof_FEC.Data[4726] := 358.11;
   Prof_FEC.Data[4727] := 307.2;
   Prof_FEC.Data[4728] := 371.53;
   Prof_FEC.Data[4729] := 387.72;
   Prof_FEC.Data[4730] := 385.93;
   Prof_FEC.Data[4731] := 374.95;
   Prof_FEC.Data[4732] := 371.68;
   Prof_FEC.Data[4733] := 421.89;
   Prof_FEC.Data[4734] := 396.51;
   Prof_FEC.Data[4735] := 447.36;
   Prof_FEC.Data[4736] := 466.5;
   Prof_FEC.Data[4737] := 478.34;
   Prof_FEC.Data[4738] := 487.98;
   Prof_FEC.Data[4739] := 505.43;
   Prof_FEC.Data[4740] := 572.99;
   Prof_FEC.Data[4741] := 573.25;
   Prof_FEC.Data[4742] := 612.06;
   Prof_FEC.Data[4743] := 663.6;
   Prof_FEC.Data[4744] := 639.31;
   Prof_FEC.Data[4745] := 660.8;
   Prof_FEC.Data[4746] := 698.77;
   Prof_FEC.Data[4747] := 575.52;
   Prof_FEC.Data[4748] := 620.6;
   Prof_FEC.Data[4749] := 662.5;
   Prof_FEC.Data[4750] := 633.41;
   Prof_FEC.Data[4751] := 668.79;
   Prof_FEC.Data[4752] := 634.65;
   Prof_FEC.Data[4753] := 575.77;
   Prof_FEC.Data[4754] := 550.11;
   Prof_FEC.Data[4755] := 577.32;
   Prof_FEC.Data[4756] := 549.15;
   Prof_FEC.Data[4757] := 711.43;
   Prof_FEC.Data[4758] := 675.1;
   Prof_FEC.Data[4759] := 605.85;
   Prof_FEC.Data[4760] := 526.06;
   Prof_FEC.Data[4761] := 584.7;
   Prof_FEC.Data[4762] := 534.19;
   Prof_FEC.Data[4763] := 577.53;
   Prof_FEC.Data[4764] := 518.77;
   Prof_FEC.Data[4765] := 657.33;
   Prof_FEC.Data[4766] := 611.33;
   Prof_FEC.Data[4767] := 557.98;
   Prof_FEC.Data[4768] := 672.26;
   Prof_FEC.Data[4769] := 667.22;
   Prof_FEC.Data[4770] := 620.59;
   Prof_FEC.Data[4771] := 594.79;
   Prof_FEC.Data[4772] := 394.39;
   Prof_FEC.Data[4773] := 352.02;
   Prof_FEC.Data[4774] := 292.57;
   Prof_FEC.Data[4775] := 297.29;
   Prof_FEC.Data[4776] := 256.77;
   Prof_FEC.Data[4777] := 253.38;
   Prof_FEC.Data[4778] := 226.58;
   Prof_FEC.Data[4779] := 263.13;
   Prof_FEC.Data[4780] := 42.591;
   Prof_FEC.Data[4781] := 43.786;
   Prof_FEC.Data[4782] := 42.501;
   Prof_FEC.Data[4783] := 43.203;
   Prof_FEC.Data[4784] := 37.248;
   Prof_FEC.Data[4785] := 38.5;
   Prof_FEC.Data[4786] := 37.164;
   Prof_FEC.Data[4787] := 37.842;
   Prof_FEC.Data[4788] := 41.036;
   Prof_FEC.Data[4789] := 46.165;
   Prof_FEC.Data[4790] := 44.022;
   Prof_FEC.Data[4791] := 43.434;
   Prof_FEC.Data[4792] := 42.865;
   Prof_FEC.Data[4793] := 40.073;
   Prof_FEC.Data[4794] := 42.062;
   Prof_FEC.Data[4795] := 42.304;
   Prof_FEC.Data[4796] := 45.346;
   Prof_FEC.Data[4797] := 43.944;
   Prof_FEC.Data[4798] := 46.085;
   Prof_FEC.Data[4799] := 41.492;
   Prof_FEC.Data[4800] := 42.46;
   Prof_FEC.Data[4801] := 43.692;
   Prof_FEC.Data[4802] := 42.376;
   Prof_FEC.Data[4803] := 43.761;
   Prof_FEC.Data[4804] := 50.0;
   Prof_FEC.Data[4805] := 50.0;
   Prof_FEC.Data[4806] := 47.188;
   Prof_FEC.Data[4807] := 44.145;
   Prof_FEC.Data[4808] := 39.92;
   Prof_FEC.Data[4809] := 43.558;
   Prof_FEC.Data[4810] := 44.397;
   Prof_FEC.Data[4811] := 42.712;
   Prof_FEC.Data[4812] := 41.55;
   Prof_FEC.Data[4813] := 43.586;
   Prof_FEC.Data[4814] := 42.725;
   Prof_FEC.Data[4815] := 41.657;
   Prof_FEC.Data[4816] := 42.875;
   Prof_FEC.Data[4817] := 41.164;
   Prof_FEC.Data[4818] := 42.509;
   Prof_FEC.Data[4819] := 42.977;
   Prof_FEC.Data[4820] := 282.36;
   Prof_FEC.Data[4821] := 279.35;
   Prof_FEC.Data[4822] := 300.6;
   Prof_FEC.Data[4823] := 305.94;
   Prof_FEC.Data[4824] := 343.07;
   Prof_FEC.Data[4825] := 375.64;
   Prof_FEC.Data[4826] := 333.97;
   Prof_FEC.Data[4827] := 369.84;
   Prof_FEC.Data[4828] := 396.77;
   Prof_FEC.Data[4829] := 410.41;
   Prof_FEC.Data[4830] := 423.43;
   Prof_FEC.Data[4831] := 426.92;
   Prof_FEC.Data[4832] := 509.23;
   Prof_FEC.Data[4833] := 549.89;
   Prof_FEC.Data[4834] := 599.89;
   Prof_FEC.Data[4835] := 599.75;
   Prof_FEC.Data[4836] := 601.55;
   Prof_FEC.Data[4837] := 606.68;
   Prof_FEC.Data[4838] := 595.03;
   Prof_FEC.Data[4839] := 638.44;
   Prof_FEC.Data[4840] := 650.5;
   Prof_FEC.Data[4841] := 677.58;
   Prof_FEC.Data[4842] := 626.45;
   Prof_FEC.Data[4843] := 667.22;
   Prof_FEC.Data[4844] := 636.54;
   Prof_FEC.Data[4845] := 640.55;
   Prof_FEC.Data[4846] := 724.58;
   Prof_FEC.Data[4847] := 676.71;
   Prof_FEC.Data[4848] := 631.45;
   Prof_FEC.Data[4849] := 612.06;
   Prof_FEC.Data[4850] := 662.98;
   Prof_FEC.Data[4851] := 664.84;
   Prof_FEC.Data[4852] := 736.05;
   Prof_FEC.Data[4853] := 700.15;
   Prof_FEC.Data[4854] := 678.3;
   Prof_FEC.Data[4855] := 694.37;
   Prof_FEC.Data[4856] := 769.14;
   Prof_FEC.Data[4857] := 706.03;
   Prof_FEC.Data[4858] := 717.17;
   Prof_FEC.Data[4859] := 775.21;
   Prof_FEC.Data[4860] := 711.64;
   Prof_FEC.Data[4861] := 701.63;
   Prof_FEC.Data[4862] := 673.17;
   Prof_FEC.Data[4863] := 741.17;
   Prof_FEC.Data[4864] := 743.99;
   Prof_FEC.Data[4865] := 709.08;
   Prof_FEC.Data[4866] := 687.13;
   Prof_FEC.Data[4867] := 624.5;
   Prof_FEC.Data[4868] := 404.65;
   Prof_FEC.Data[4869] := 321.3;
   Prof_FEC.Data[4870] := 315.45;
   Prof_FEC.Data[4871] := 277.86;
   Prof_FEC.Data[4872] := 266.5;
   Prof_FEC.Data[4873] := 252.12;
   Prof_FEC.Data[4874] := 281.85;
   Prof_FEC.Data[4875] := 273.29;
   Prof_FEC.Data[4876] := 42.448;
   Prof_FEC.Data[4877] := 43.289;
   Prof_FEC.Data[4878] := 42.637;
   Prof_FEC.Data[4879] := 38.596;
   Prof_FEC.Data[4880] := 36.78;
   Prof_FEC.Data[4881] := 36.083;
   Prof_FEC.Data[4882] := 35.672;
   Prof_FEC.Data[4883] := 38.067;
   Prof_FEC.Data[4884] := 37.359;
   Prof_FEC.Data[4885] := 40.19;
   Prof_FEC.Data[4886] := 39.351;
   Prof_FEC.Data[4887] := 40.138;
   Prof_FEC.Data[4888] := 36.497;
   Prof_FEC.Data[4889] := 39.197;
   Prof_FEC.Data[4890] := 38.142;
   Prof_FEC.Data[4891] := 39.915;
   Prof_FEC.Data[4892] := 41.446;
   Prof_FEC.Data[4893] := 41.984;
   Prof_FEC.Data[4894] := 40.728;
   Prof_FEC.Data[4895] := 41.215;
   Prof_FEC.Data[4896] := 38.314;
   Prof_FEC.Data[4897] := 37.091;
   Prof_FEC.Data[4898] := 39.908;
   Prof_FEC.Data[4899] := 42.239;
   Prof_FEC.Data[4900] := 41.238;
   Prof_FEC.Data[4901] := 43.221;
   Prof_FEC.Data[4902] := 43.532;
   Prof_FEC.Data[4903] := 40.226;
   Prof_FEC.Data[4904] := 38.465;
   Prof_FEC.Data[4905] := 39.579;
   Prof_FEC.Data[4906] := 39.024;
   Prof_FEC.Data[4907] := 39.725;
   Prof_FEC.Data[4908] := 40.784;
   Prof_FEC.Data[4909] := 41.632;
   Prof_FEC.Data[4910] := 41.086;
   Prof_FEC.Data[4911] := 40.968;
   Prof_FEC.Data[4912] := 38.803;
   Prof_FEC.Data[4913] := 40.215;
   Prof_FEC.Data[4914] := 39.961;
   Prof_FEC.Data[4915] := 41.824;
   Prof_FEC.Data[4916] := 275.0;
   Prof_FEC.Data[4917] := 259.61;
   Prof_FEC.Data[4918] := 262.0;
   Prof_FEC.Data[4919] := 337.73;
   Prof_FEC.Data[4920] := 380.06;
   Prof_FEC.Data[4921] := 385.88;
   Prof_FEC.Data[4922] := 423.79;
   Prof_FEC.Data[4923] := 410.1;
   Prof_FEC.Data[4924] := 434.41;
   Prof_FEC.Data[4925] := 444.69;
   Prof_FEC.Data[4926] := 443.53;
   Prof_FEC.Data[4927] := 480.63;
   Prof_FEC.Data[4928] := 507.36;
   Prof_FEC.Data[4929] := 539.64;
   Prof_FEC.Data[4930] := 547.46;
   Prof_FEC.Data[4931] := 575.06;
   Prof_FEC.Data[4932] := 584.2;
   Prof_FEC.Data[4933] := 616.65;
   Prof_FEC.Data[4934] := 676.31;
   Prof_FEC.Data[4935] := 666.19;
   Prof_FEC.Data[4936] := 566.23;
   Prof_FEC.Data[4937] := 579.03;
   Prof_FEC.Data[4938] := 693.28;
   Prof_FEC.Data[4939] := 684.17;
   Prof_FEC.Data[4940] := 631.46;
   Prof_FEC.Data[4941] := 686.47;
   Prof_FEC.Data[4942] := 702.42;
   Prof_FEC.Data[4943] := 663.74;
   Prof_FEC.Data[4944] := 677.03;
   Prof_FEC.Data[4945] := 596.34;
   Prof_FEC.Data[4946] := 657.12;
   Prof_FEC.Data[4947] := 643.2;
   Prof_FEC.Data[4948] := 631.68;
   Prof_FEC.Data[4949] := 675.17;
   Prof_FEC.Data[4950] := 642.06;
   Prof_FEC.Data[4951] := 633.67;
   Prof_FEC.Data[4952] := 654.81;
   Prof_FEC.Data[4953] := 633.42;
   Prof_FEC.Data[4954] := 669.17;
   Prof_FEC.Data[4955] := 672.16;
   Prof_FEC.Data[4956] := 773.03;
   Prof_FEC.Data[4957] := 652.47;
   Prof_FEC.Data[4958] := 802.85;
   Prof_FEC.Data[4959] := 685.87;
   Prof_FEC.Data[4960] := 787.95;
   Prof_FEC.Data[4961] := 715.39;
   Prof_FEC.Data[4962] := 602.25;
   Prof_FEC.Data[4963] := 574.13;
   Prof_FEC.Data[4964] := 375.57;
   Prof_FEC.Data[4965] := 321.37;
   Prof_FEC.Data[4966] := 273.01;
   Prof_FEC.Data[4967] := 261.13;
   Prof_FEC.Data[4968] := 256.13;
   Prof_FEC.Data[4969] := 251.5;
   Prof_FEC.Data[4970] := 234.48;
   Prof_FEC.Data[4971] := 251.15;
   Prof_FEC.Data[4972] := 43.535;
   Prof_FEC.Data[4973] := 43.089;
   Prof_FEC.Data[4974] := 41.617;
   Prof_FEC.Data[4975] := 42.784;
   Prof_FEC.Data[4976] := 40.007;
   Prof_FEC.Data[4977] := 42.897;
   Prof_FEC.Data[4978] := 43.2;
   Prof_FEC.Data[4979] := 42.191;
   Prof_FEC.Data[4980] := 45.753;
   Prof_FEC.Data[4981] := 48.353;
   Prof_FEC.Data[4982] := 44.436;
   Prof_FEC.Data[4983] := 46.377;
   Prof_FEC.Data[4984] := 43.505;
   Prof_FEC.Data[4985] := 45.634;
   Prof_FEC.Data[4986] := 44.013;
   Prof_FEC.Data[4987] := 44.408;
   Prof_FEC.Data[4988] := 46.66;
   Prof_FEC.Data[4989] := 46.125;
   Prof_FEC.Data[4990] := 45.22;
   Prof_FEC.Data[4991] := 46.536;
   Prof_FEC.Data[4992] := 42.58;
   Prof_FEC.Data[4993] := 41.82;
   Prof_FEC.Data[4994] := 42.289;
   Prof_FEC.Data[4995] := 44.775;
   Prof_FEC.Data[4996] := 46.98;
   Prof_FEC.Data[4997] := 46.934;
   Prof_FEC.Data[4998] := 43.384;
   Prof_FEC.Data[4999] := 48.065;
   Prof_FEC.Data[5000] := 41.714;
   Prof_FEC.Data[5001] := 39.813;
   Prof_FEC.Data[5002] := 41.216;
   Prof_FEC.Data[5003] := 45.705;
   Prof_FEC.Data[5004] := 46.942;
   Prof_FEC.Data[5005] := 46.718;
   Prof_FEC.Data[5006] := 44.278;
   Prof_FEC.Data[5007] := 44.62;
   Prof_FEC.Data[5008] := 45.625;
   Prof_FEC.Data[5009] := 42.933;
   Prof_FEC.Data[5010] := 43.246;
   Prof_FEC.Data[5011] := 43.895;
   Prof_FEC.Data[5012] := 320.63;
   Prof_FEC.Data[5013] := 309.86;
   Prof_FEC.Data[5014] := 271.77;
   Prof_FEC.Data[5015] := 276.65;
   Prof_FEC.Data[5016] := 232.53;
   Prof_FEC.Data[5017] := 213.78;
   Prof_FEC.Data[5018] := 224.63;
   Prof_FEC.Data[5019] := 232.19;
   Prof_FEC.Data[5020] := 215.79;
   Prof_FEC.Data[5021] := 223.78;
   Prof_FEC.Data[5022] := 214.17;
   Prof_FEC.Data[5023] := 221.94;
   Prof_FEC.Data[5024] := 242.28;
   Prof_FEC.Data[5025] := 250.25;
   Prof_FEC.Data[5026] := 267.21;
   Prof_FEC.Data[5027] := 278.76;
   Prof_FEC.Data[5028] := 281.35;
   Prof_FEC.Data[5029] := 302.33;
   Prof_FEC.Data[5030] := 325.65;
   Prof_FEC.Data[5031] := 342.05;
   Prof_FEC.Data[5032] := 311.73;
   Prof_FEC.Data[5033] := 300.4;
   Prof_FEC.Data[5034] := 341.78;
   Prof_FEC.Data[5035] := 317.26;
   Prof_FEC.Data[5036] := 327.11;
   Prof_FEC.Data[5037] := 349.58;
   Prof_FEC.Data[5038] := 338.6;
   Prof_FEC.Data[5039] := 312.0;
   Prof_FEC.Data[5040] := 274.98;
   Prof_FEC.Data[5041] := 246.24;
   Prof_FEC.Data[5042] := 239.54;
   Prof_FEC.Data[5043] := 239.98;
   Prof_FEC.Data[5044] := 208.94;
   Prof_FEC.Data[5045] := 251.5;
   Prof_FEC.Data[5046] := 227.2;
   Prof_FEC.Data[5047] := 230.02;
   Prof_FEC.Data[5048] := 282.75;
   Prof_FEC.Data[5049] := 285.58;
   Prof_FEC.Data[5050] := 290.67;
   Prof_FEC.Data[5051] := 271.79;
   Prof_FEC.Data[5052] := 323.12;
   Prof_FEC.Data[5053] := 319.08;
   Prof_FEC.Data[5054] := 275.63;
   Prof_FEC.Data[5055] := 250.83;
   Prof_FEC.Data[5056] := 178.79;
   Prof_FEC.Data[5057] := 137.07;
   Prof_FEC.Data[5058] := 121.03;
   Prof_FEC.Data[5059] := 149.01;
   Prof_FEC.Data[5060] := 171.04;
   Prof_FEC.Data[5061] := 169.36;
   Prof_FEC.Data[5062] := 192.12;
   Prof_FEC.Data[5063] := 193.02;
   Prof_FEC.Data[5064] := 267.47;
   Prof_FEC.Data[5065] := 294.39;
   Prof_FEC.Data[5066] := 276.56;
   Prof_FEC.Data[5067] := 276.24;
   Prof_FEC.Data[5068] := 39.313;
   Prof_FEC.Data[5069] := 40.0;
   Prof_FEC.Data[5070] := 38.275;
   Prof_FEC.Data[5071] := 40.226;
   Prof_FEC.Data[5072] := 40.947;
   Prof_FEC.Data[5073] := 43.36;
   Prof_FEC.Data[5074] := 41.77;
   Prof_FEC.Data[5075] := 45.318;
   Prof_FEC.Data[5076] := 40.96;
   Prof_FEC.Data[5077] := 39.276;
   Prof_FEC.Data[5078] := 43.171;
   Prof_FEC.Data[5079] := 38.79;
   Prof_FEC.Data[5080] := 43.118;
   Prof_FEC.Data[5081] := 42.188;
   Prof_FEC.Data[5082] := 43.063;
   Prof_FEC.Data[5083] := 42.18;
   Prof_FEC.Data[5084] := 44.761;
   Prof_FEC.Data[5085] := 41.131;
   Prof_FEC.Data[5086] := 41.051;
   Prof_FEC.Data[5087] := 43.515;
   Prof_FEC.Data[5088] := 45.604;
   Prof_FEC.Data[5089] := 46.753;
   Prof_FEC.Data[5090] := 48.248;
   Prof_FEC.Data[5091] := 47.625;
   Prof_FEC.Data[5092] := 40.785;
   Prof_FEC.Data[5093] := 42.852;
   Prof_FEC.Data[5094] := 42.167;
   Prof_FEC.Data[5095] := 42.466;
   Prof_FEC.Data[5096] := 43.503;
   Prof_FEC.Data[5097] := 44.685;
   Prof_FEC.Data[5098] := 44.29;
   Prof_FEC.Data[5099] := 47.765;
   Prof_FEC.Data[5100] := 42.796;
   Prof_FEC.Data[5101] := 40.122;
   Prof_FEC.Data[5102] := 43.293;
   Prof_FEC.Data[5103] := 42.252;
   Prof_FEC.Data[5104] := 43.065;
   Prof_FEC.Data[5105] := 44.049;
   Prof_FEC.Data[5106] := 43.032;
   Prof_FEC.Data[5107] := 41.792;
   Prof_FEC.Data[5108] := 255.03;
   Prof_FEC.Data[5109] := 272.98;
   Prof_FEC.Data[5110] := 244.05;
   Prof_FEC.Data[5111] := 266.94;
   Prof_FEC.Data[5112] := 277.22;
   Prof_FEC.Data[5113] := 306.35;
   Prof_FEC.Data[5114] := 260.72;
   Prof_FEC.Data[5115] := 257.08;
   Prof_FEC.Data[5116] := 199.05;
   Prof_FEC.Data[5117] := 159.25;
   Prof_FEC.Data[5118] := 151.14;
   Prof_FEC.Data[5119] := 138.94;
   Prof_FEC.Data[5120] := 160.47;
   Prof_FEC.Data[5121] := 170.1;
   Prof_FEC.Data[5122] := 166.62;
   Prof_FEC.Data[5123] := 167.5;
   Prof_FEC.Data[5124] := 146.17;
   Prof_FEC.Data[5125] := 132.5;
   Prof_FEC.Data[5126] := 143.29;
   Prof_FEC.Data[5127] := 141.95;
   Prof_FEC.Data[5128] := 145.02;
   Prof_FEC.Data[5129] := 150.1;
   Prof_FEC.Data[5130] := 157.37;
   Prof_FEC.Data[5131] := 149.13;
   Prof_FEC.Data[5132] := 109.86;
   Prof_FEC.Data[5133] := 106.81;
   Prof_FEC.Data[5134] := 111.08;
   Prof_FEC.Data[5135] := 110.15;
   Prof_FEC.Data[5136] := 127.03;
   Prof_FEC.Data[5137] := 132.4;
   Prof_FEC.Data[5138] := 135.7;
   Prof_FEC.Data[5139] := 128.33;
   Prof_FEC.Data[5140] := 109.69;
   Prof_FEC.Data[5141] := 114.98;
   Prof_FEC.Data[5142] := 103.0;
   Prof_FEC.Data[5143] := 121.89;
   Prof_FEC.Data[5144] := 137.41;
   Prof_FEC.Data[5145] := 138.79;
   Prof_FEC.Data[5146] := 134.6;
   Prof_FEC.Data[5147] := 148.62;
   Prof_FEC.Data[5148] := 135.69;
   Prof_FEC.Data[5149] := 137.92;
   Prof_FEC.Data[5150] := 134.61;
   Prof_FEC.Data[5151] := 118.35;
   Prof_FEC.Data[5152] := 136.23;
   Prof_FEC.Data[5153] := 137.91;
   Prof_FEC.Data[5154] := 151.31;
   Prof_FEC.Data[5155] := 152.69;
   Prof_FEC.Data[5156] := 163.02;
   Prof_FEC.Data[5157] := 180.6;
   Prof_FEC.Data[5158] := 181.65;
   Prof_FEC.Data[5159] := 202.16;
   Prof_FEC.Data[5160] := 257.91;
   Prof_FEC.Data[5161] := 243.22;
   Prof_FEC.Data[5162] := 289.31;
   Prof_FEC.Data[5163] := 251.26;
   Prof_FEC.Data[5164] := 38.809;
   Prof_FEC.Data[5165] := 39.735;
   Prof_FEC.Data[5166] := 37.666;
   Prof_FEC.Data[5167] := 38.589;
   Prof_FEC.Data[5168] := 43.571;
   Prof_FEC.Data[5169] := 39.438;
   Prof_FEC.Data[5170] := 44.345;
   Prof_FEC.Data[5171] := 40.563;
   Prof_FEC.Data[5172] := 39.691;
   Prof_FEC.Data[5173] := 41.563;
   Prof_FEC.Data[5174] := 36.695;
   Prof_FEC.Data[5175] := 37.525;
   Prof_FEC.Data[5176] := 40.106;
   Prof_FEC.Data[5177] := 39.34;
   Prof_FEC.Data[5178] := 41.478;
   Prof_FEC.Data[5179] := 43.274;
   Prof_FEC.Data[5180] := 40.281;
   Prof_FEC.Data[5181] := 40.819;
   Prof_FEC.Data[5182] := 39.047;
   Prof_FEC.Data[5183] := 38.618;
   Prof_FEC.Data[5184] := 41.754;
   Prof_FEC.Data[5185] := 39.791;
   Prof_FEC.Data[5186] := 41.722;
   Prof_FEC.Data[5187] := 41.831;
   Prof_FEC.Data[5188] := 38.778;
   Prof_FEC.Data[5189] := 40.578;
   Prof_FEC.Data[5190] := 41.218;
   Prof_FEC.Data[5191] := 40.62;
   Prof_FEC.Data[5192] := 43.504;
   Prof_FEC.Data[5193] := 40.86;
   Prof_FEC.Data[5194] := 41.376;
   Prof_FEC.Data[5195] := 43.896;
   Prof_FEC.Data[5196] := 43.706;
   Prof_FEC.Data[5197] := 41.155;
   Prof_FEC.Data[5198] := 41.083;
   Prof_FEC.Data[5199] := 38.464;
   Prof_FEC.Data[5200] := 41.771;
   Prof_FEC.Data[5201] := 43.332;
   Prof_FEC.Data[5202] := 45.483;
   Prof_FEC.Data[5203] := 42.442;
   Prof_FEC.Data[5204] := 259.17;
   Prof_FEC.Data[5205] := 225.36;
   Prof_FEC.Data[5206] := 258.48;
   Prof_FEC.Data[5207] := 242.98;
   Prof_FEC.Data[5208] := 291.23;
   Prof_FEC.Data[5209] := 298.74;
   Prof_FEC.Data[5210] := 265.63;
   Prof_FEC.Data[5211] := 227.71;
   Prof_FEC.Data[5212] := 189.26;
   Prof_FEC.Data[5213] := 147.48;
   Prof_FEC.Data[5214] := 131.6;
   Prof_FEC.Data[5215] := 128.57;
   Prof_FEC.Data[5216] := 147.95;
   Prof_FEC.Data[5217] := 141.66;
   Prof_FEC.Data[5218] := 132.08;
   Prof_FEC.Data[5219] := 117.24;
   Prof_FEC.Data[5220] := 99.44;
   Prof_FEC.Data[5221] := 98.52;
   Prof_FEC.Data[5222] := 99.86;
   Prof_FEC.Data[5223] := 112.24;
   Prof_FEC.Data[5224] := 117.79;
   Prof_FEC.Data[5225] := 139.2;
   Prof_FEC.Data[5226] := 119.86;
   Prof_FEC.Data[5227] := 111.72;
   Prof_FEC.Data[5228] := 97.75;
   Prof_FEC.Data[5229] := 113.64;
   Prof_FEC.Data[5230] := 98.32;
   Prof_FEC.Data[5231] := 108.43;
   Prof_FEC.Data[5232] := 128.62;
   Prof_FEC.Data[5233] := 129.17;
   Prof_FEC.Data[5234] := 122.14;
   Prof_FEC.Data[5235] := 117.45;
   Prof_FEC.Data[5236] := 114.95;
   Prof_FEC.Data[5237] := 105.79;
   Prof_FEC.Data[5238] := 112.54;
   Prof_FEC.Data[5239] := 114.69;
   Prof_FEC.Data[5240] := 122.15;
   Prof_FEC.Data[5241] := 113.55;
   Prof_FEC.Data[5242] := 117.57;
   Prof_FEC.Data[5243] := 100.63;
   Prof_FEC.Data[5244] := 95.62;
   Prof_FEC.Data[5245] := 94.67;
   Prof_FEC.Data[5246] := 106.4;
   Prof_FEC.Data[5247] := 110.82;
   Prof_FEC.Data[5248] := 101.74;
   Prof_FEC.Data[5249] := 102.63;
   Prof_FEC.Data[5250] := 106.67;
   Prof_FEC.Data[5251] := 119.67;
   Prof_FEC.Data[5252] := 154.66;
   Prof_FEC.Data[5253] := 160.55;
   Prof_FEC.Data[5254] := 170.61;
   Prof_FEC.Data[5255] := 193.96;
   Prof_FEC.Data[5256] := 199.09;
   Prof_FEC.Data[5257] := 212.69;
   Prof_FEC.Data[5258] := 229.18;
   Prof_FEC.Data[5259] := 207.73;
   Prof_FEC.Data[5260] := 34.656;
   Prof_FEC.Data[5261] := 35.367;
   Prof_FEC.Data[5262] := 38.156;
   Prof_FEC.Data[5263] := 36.193;
   Prof_FEC.Data[5264] := 37.556;
   Prof_FEC.Data[5265] := 36.735;
   Prof_FEC.Data[5266] := 38.079;
   Prof_FEC.Data[5267] := 36.984;
   Prof_FEC.Data[5268] := 37.407;
   Prof_FEC.Data[5269] := 35.969;
   Prof_FEC.Data[5270] := 37.329;
   Prof_FEC.Data[5271] := 37.688;
   Prof_FEC.Data[5272] := 38.992;
   Prof_FEC.Data[5273] := 39.958;
   Prof_FEC.Data[5274] := 40.654;
   Prof_FEC.Data[5275] := 39.448;
   Prof_FEC.Data[5276] := 36.842;
   Prof_FEC.Data[5277] := 36.444;
   Prof_FEC.Data[5278] := 36.304;
   Prof_FEC.Data[5279] := 37.053;
   Prof_FEC.Data[5280] := 37.917;
   Prof_FEC.Data[5281] := 38.311;
   Prof_FEC.Data[5282] := 39.706;
   Prof_FEC.Data[5283] := 39.724;
   Prof_FEC.Data[5284] := 35.065;
   Prof_FEC.Data[5285] := 34.985;
   Prof_FEC.Data[5286] := 35.846;
   Prof_FEC.Data[5287] := 36.904;
   Prof_FEC.Data[5288] := 37.143;
   Prof_FEC.Data[5289] := 41.588;
   Prof_FEC.Data[5290] := 41.174;
   Prof_FEC.Data[5291] := 37.465;
   Prof_FEC.Data[5292] := 37.494;
   Prof_FEC.Data[5293] := 37.967;
   Prof_FEC.Data[5294] := 35.801;
   Prof_FEC.Data[5295] := 39.504;
   Prof_FEC.Data[5296] := 39.894;
   Prof_FEC.Data[5297] := 39.984;
   Prof_FEC.Data[5298] := 38.894;
   Prof_FEC.Data[5299] := 40.273;
   Prof_FEC.Data[5300] := 196.36;
   Prof_FEC.Data[5301] := 198.55;
   Prof_FEC.Data[5302] := 224.92;
   Prof_FEC.Data[5303] := 267.63;
   Prof_FEC.Data[5304] := 367.66;
   Prof_FEC.Data[5305] := 412.7;
   Prof_FEC.Data[5306] := 429.4;
   Prof_FEC.Data[5307] := 446.79;
   Prof_FEC.Data[5308] := 407.5;
   Prof_FEC.Data[5309] := 411.2;
   Prof_FEC.Data[5310] := 475.94;
   Prof_FEC.Data[5311] := 479.92;
   Prof_FEC.Data[5312] := 564.14;
   Prof_FEC.Data[5313] := 621.22;
   Prof_FEC.Data[5314] := 656.26;
   Prof_FEC.Data[5315] := 650.73;
   Prof_FEC.Data[5316] := 692.74;
   Prof_FEC.Data[5317] := 710.87;
   Prof_FEC.Data[5318] := 743.97;
   Prof_FEC.Data[5319] := 760.46;
   Prof_FEC.Data[5320] := 737.02;
   Prof_FEC.Data[5321] := 684.35;
   Prof_FEC.Data[5322] := 725.88;
   Prof_FEC.Data[5323] := 663.61;
   Prof_FEC.Data[5324] := 643.39;
   Prof_FEC.Data[5325] := 652.68;
   Prof_FEC.Data[5326] := 650.79;
   Prof_FEC.Data[5327] := 609.53;
   Prof_FEC.Data[5328] := 614.76;
   Prof_FEC.Data[5329] := 650.47;
   Prof_FEC.Data[5330] := 594.67;
   Prof_FEC.Data[5331] := 658.21;
   Prof_FEC.Data[5332] := 596.13;
   Prof_FEC.Data[5333] := 713.16;
   Prof_FEC.Data[5334] := 737.91;
   Prof_FEC.Data[5335] := 776.67;
   Prof_FEC.Data[5336] := 753.95;
   Prof_FEC.Data[5337] := 694.69;
   Prof_FEC.Data[5338] := 655.1;
   Prof_FEC.Data[5339] := 693.35;
   Prof_FEC.Data[5340] := 686.84;
   Prof_FEC.Data[5341] := 723.97;
   Prof_FEC.Data[5342] := 655.1;
   Prof_FEC.Data[5343] := 651.49;
   Prof_FEC.Data[5344] := 669.85;
   Prof_FEC.Data[5345] := 671.68;
   Prof_FEC.Data[5346] := 679.04;
   Prof_FEC.Data[5347] := 556.55;
   Prof_FEC.Data[5348] := 310.55;
   Prof_FEC.Data[5349] := 251.93;
   Prof_FEC.Data[5350] := 223.74;
   Prof_FEC.Data[5351] := 203.14;
   Prof_FEC.Data[5352] := 211.53;
   Prof_FEC.Data[5353] := 215.71;
   Prof_FEC.Data[5354] := 189.66;
   Prof_FEC.Data[5355] := 193.7;
   Prof_FEC.Data[5356] := 38.348;
   Prof_FEC.Data[5357] := 35.497;
   Prof_FEC.Data[5358] := 36.598;
   Prof_FEC.Data[5359] := 34.475;
   Prof_FEC.Data[5360] := 34.415;
   Prof_FEC.Data[5361] := 33.754;
   Prof_FEC.Data[5362] := 34.461;
   Prof_FEC.Data[5363] := 36.181;
   Prof_FEC.Data[5364] := 38.887;
   Prof_FEC.Data[5365] := 38.879;
   Prof_FEC.Data[5366] := 39.241;
   Prof_FEC.Data[5367] := 38.65;
   Prof_FEC.Data[5368] := 34.676;
   Prof_FEC.Data[5369] := 37.533;
   Prof_FEC.Data[5370] := 36.361;
   Prof_FEC.Data[5371] := 38.372;
   Prof_FEC.Data[5372] := 36.379;
   Prof_FEC.Data[5373] := 39.898;
   Prof_FEC.Data[5374] := 39.957;
   Prof_FEC.Data[5375] := 39.52;
   Prof_FEC.Data[5376] := 37.135;
   Prof_FEC.Data[5377] := 36.687;
   Prof_FEC.Data[5378] := 36.698;
   Prof_FEC.Data[5379] := 38.255;
   Prof_FEC.Data[5380] := 40.449;
   Prof_FEC.Data[5381] := 39.906;
   Prof_FEC.Data[5382] := 40.131;
   Prof_FEC.Data[5383] := 37.944;
   Prof_FEC.Data[5384] := 39.318;
   Prof_FEC.Data[5385] := 37.693;
   Prof_FEC.Data[5386] := 36.221;
   Prof_FEC.Data[5387] := 39.475;
   Prof_FEC.Data[5388] := 39.897;
   Prof_FEC.Data[5389] := 38.273;
   Prof_FEC.Data[5390] := 39.196;
   Prof_FEC.Data[5391] := 37.848;
   Prof_FEC.Data[5392] := 34.85;
   Prof_FEC.Data[5393] := 37.857;
   Prof_FEC.Data[5394] := 36.553;
   Prof_FEC.Data[5395] := 40.682;
   Prof_FEC.Data[5396] := 198.86;
   Prof_FEC.Data[5397] := 199.04;
   Prof_FEC.Data[5398] := 268.65;
   Prof_FEC.Data[5399] := 274.39;
   Prof_FEC.Data[5400] := 333.42;
   Prof_FEC.Data[5401] := 366.9;
   Prof_FEC.Data[5402] := 338.43;
   Prof_FEC.Data[5403] := 343.66;
   Prof_FEC.Data[5404] := 404.44;
   Prof_FEC.Data[5405] := 356.2;
   Prof_FEC.Data[5406] := 440.67;
   Prof_FEC.Data[5407] := 436.06;
   Prof_FEC.Data[5408] := 476.46;
   Prof_FEC.Data[5409] := 448.72;
   Prof_FEC.Data[5410] := 559.64;
   Prof_FEC.Data[5411] := 492.31;
   Prof_FEC.Data[5412] := 536.11;
   Prof_FEC.Data[5413] := 565.24;
   Prof_FEC.Data[5414] := 562.74;
   Prof_FEC.Data[5415] := 575.05;
   Prof_FEC.Data[5416] := 627.62;
   Prof_FEC.Data[5417] := 653.09;
   Prof_FEC.Data[5418] := 715.1;
   Prof_FEC.Data[5419] := 691.66;
   Prof_FEC.Data[5420] := 586.87;
   Prof_FEC.Data[5421] := 665.95;
   Prof_FEC.Data[5422] := 561.8;
   Prof_FEC.Data[5423] := 535.36;
   Prof_FEC.Data[5424] := 529.27;
   Prof_FEC.Data[5425] := 507.21;
   Prof_FEC.Data[5426] := 506.43;
   Prof_FEC.Data[5427] := 447.71;
   Prof_FEC.Data[5428] := 555.63;
   Prof_FEC.Data[5429] := 587.03;
   Prof_FEC.Data[5430] := 588.66;
   Prof_FEC.Data[5431] := 541.09;
   Prof_FEC.Data[5432] := 615.54;
   Prof_FEC.Data[5433] := 600.3;
   Prof_FEC.Data[5434] := 596.36;
   Prof_FEC.Data[5435] := 567.5;
   Prof_FEC.Data[5436] := 665.05;
   Prof_FEC.Data[5437] := 621.98;
   Prof_FEC.Data[5438] := 643.45;
   Prof_FEC.Data[5439] := 640.5;
   Prof_FEC.Data[5440] := 701.37;
   Prof_FEC.Data[5441] := 678.74;
   Prof_FEC.Data[5442] := 614.59;
   Prof_FEC.Data[5443] := 541.84;
   Prof_FEC.Data[5444] := 345.93;
   Prof_FEC.Data[5445] := 280.46;
   Prof_FEC.Data[5446] := 196.25;
   Prof_FEC.Data[5447] := 211.45;
   Prof_FEC.Data[5448] := 194.98;
   Prof_FEC.Data[5449] := 218.14;
   Prof_FEC.Data[5450] := 184.36;
   Prof_FEC.Data[5451] := 212.17;
   Prof_FEC.Data[5452] := 38.581;
   Prof_FEC.Data[5453] := 38.621;
   Prof_FEC.Data[5454] := 38.166;
   Prof_FEC.Data[5455] := 37.894;
   Prof_FEC.Data[5456] := 37.963;
   Prof_FEC.Data[5457] := 39.208;
   Prof_FEC.Data[5458] := 38.739;
   Prof_FEC.Data[5459] := 36.763;
   Prof_FEC.Data[5460] := 41.508;
   Prof_FEC.Data[5461] := 41.803;
   Prof_FEC.Data[5462] := 41.429;
   Prof_FEC.Data[5463] := 39.475;
   Prof_FEC.Data[5464] := 37.27;
   Prof_FEC.Data[5465] := 36.922;
   Prof_FEC.Data[5466] := 38.12;
   Prof_FEC.Data[5467] := 36.075;
   Prof_FEC.Data[5468] := 40.255;
   Prof_FEC.Data[5469] := 41.193;
   Prof_FEC.Data[5470] := 41.851;
   Prof_FEC.Data[5471] := 40.24;
   Prof_FEC.Data[5472] := 36.597;
   Prof_FEC.Data[5473] := 36.742;
   Prof_FEC.Data[5474] := 37.918;
   Prof_FEC.Data[5475] := 41.061;
   Prof_FEC.Data[5476] := 39.905;
   Prof_FEC.Data[5477] := 40.663;
   Prof_FEC.Data[5478] := 39.601;
   Prof_FEC.Data[5479] := 40.37;
   Prof_FEC.Data[5480] := 37.774;
   Prof_FEC.Data[5481] := 41.732;
   Prof_FEC.Data[5482] := 38.568;
   Prof_FEC.Data[5483] := 37.162;
   Prof_FEC.Data[5484] := 42.488;
   Prof_FEC.Data[5485] := 41.556;
   Prof_FEC.Data[5486] := 42.224;
   Prof_FEC.Data[5487] := 39.243;
   Prof_FEC.Data[5488] := 40.908;
   Prof_FEC.Data[5489] := 40.141;
   Prof_FEC.Data[5490] := 39.523;
   Prof_FEC.Data[5491] := 40.805;
   Prof_FEC.Data[5492] := 247.43;
   Prof_FEC.Data[5493] := 248.12;
   Prof_FEC.Data[5494] := 233.36;
   Prof_FEC.Data[5495] := 278.51;
   Prof_FEC.Data[5496] := 398.94;
   Prof_FEC.Data[5497] := 420.57;
   Prof_FEC.Data[5498] := 466.15;
   Prof_FEC.Data[5499] := 459.56;
   Prof_FEC.Data[5500] := 446.81;
   Prof_FEC.Data[5501] := 486.2;
   Prof_FEC.Data[5502] := 503.56;
   Prof_FEC.Data[5503] := 533.03;
   Prof_FEC.Data[5504] := 589.81;
   Prof_FEC.Data[5505] := 602.51;
   Prof_FEC.Data[5506] := 604.2;
   Prof_FEC.Data[5507] := 588.01;
   Prof_FEC.Data[5508] := 591.9;
   Prof_FEC.Data[5509] := 731.66;
   Prof_FEC.Data[5510] := 705.83;
   Prof_FEC.Data[5511] := 748.42;
   Prof_FEC.Data[5512] := 728.23;
   Prof_FEC.Data[5513] := 726.43;
   Prof_FEC.Data[5514] := 705.02;
   Prof_FEC.Data[5515] := 713.91;
   Prof_FEC.Data[5516] := 669.3;
   Prof_FEC.Data[5517] := 702.98;
   Prof_FEC.Data[5518] := 622.45;
   Prof_FEC.Data[5519] := 637.05;
   Prof_FEC.Data[5520] := 573.88;
   Prof_FEC.Data[5521] := 603.11;
   Prof_FEC.Data[5522] := 576.53;
   Prof_FEC.Data[5523] := 617.47;
   Prof_FEC.Data[5524] := 665.14;
   Prof_FEC.Data[5525] := 596.24;
   Prof_FEC.Data[5526] := 657.54;
   Prof_FEC.Data[5527] := 645.15;
   Prof_FEC.Data[5528] := 572.22;
   Prof_FEC.Data[5529] := 583.23;
   Prof_FEC.Data[5530] := 634.53;
   Prof_FEC.Data[5531] := 631.61;
   Prof_FEC.Data[5532] := 572.72;
   Prof_FEC.Data[5533] := 609.58;
   Prof_FEC.Data[5534] := 587.56;
   Prof_FEC.Data[5535] := 644.1;
   Prof_FEC.Data[5536] := 717.74;
   Prof_FEC.Data[5537] := 721.01;
   Prof_FEC.Data[5538] := 595.44;
   Prof_FEC.Data[5539] := 498.96;
   Prof_FEC.Data[5540] := 357.62;
   Prof_FEC.Data[5541] := 237.85;
   Prof_FEC.Data[5542] := 227.26;
   Prof_FEC.Data[5543] := 207.35;
   Prof_FEC.Data[5544] := 224.34;
   Prof_FEC.Data[5545] := 189.75;
   Prof_FEC.Data[5546] := 206.67;
   Prof_FEC.Data[5547] := 209.82;
   Prof_FEC.Data[5548] := 35.326;
   Prof_FEC.Data[5549] := 37.8;
   Prof_FEC.Data[5550] := 37.391;
   Prof_FEC.Data[5551] := 35.828;
   Prof_FEC.Data[5552] := 34.75;
   Prof_FEC.Data[5553] := 37.576;
   Prof_FEC.Data[5554] := 38.78;
   Prof_FEC.Data[5555] := 38.961;
   Prof_FEC.Data[5556] := 39.548;
   Prof_FEC.Data[5557] := 36.225;
   Prof_FEC.Data[5558] := 40.162;
   Prof_FEC.Data[5559] := 39.962;
   Prof_FEC.Data[5560] := 40.841;
   Prof_FEC.Data[5561] := 40.754;
   Prof_FEC.Data[5562] := 40.52;
   Prof_FEC.Data[5563] := 36.629;
   Prof_FEC.Data[5564] := 39.762;
   Prof_FEC.Data[5565] := 39.963;
   Prof_FEC.Data[5566] := 40.437;
   Prof_FEC.Data[5567] := 43.027;
   Prof_FEC.Data[5568] := 38.307;
   Prof_FEC.Data[5569] := 40.69;
   Prof_FEC.Data[5570] := 40.315;
   Prof_FEC.Data[5571] := 39.512;
   Prof_FEC.Data[5572] := 39.783;
   Prof_FEC.Data[5573] := 40.608;
   Prof_FEC.Data[5574] := 40.802;
   Prof_FEC.Data[5575] := 40.885;
   Prof_FEC.Data[5576] := 38.938;
   Prof_FEC.Data[5577] := 40.329;
   Prof_FEC.Data[5578] := 40.109;
   Prof_FEC.Data[5579] := 42.796;
   Prof_FEC.Data[5580] := 44.414;
   Prof_FEC.Data[5581] := 40.723;
   Prof_FEC.Data[5582] := 41.19;
   Prof_FEC.Data[5583] := 41.653;
   Prof_FEC.Data[5584] := 39.853;
   Prof_FEC.Data[5585] := 37.284;
   Prof_FEC.Data[5586] := 39.062;
   Prof_FEC.Data[5587] := 36.942;
   Prof_FEC.Data[5588] := 205.04;
   Prof_FEC.Data[5589] := 194.63;
   Prof_FEC.Data[5590] := 224.44;
   Prof_FEC.Data[5591] := 234.61;
   Prof_FEC.Data[5592] := 319.67;
   Prof_FEC.Data[5593] := 322.16;
   Prof_FEC.Data[5594] := 347.5;
   Prof_FEC.Data[5595] := 388.68;
   Prof_FEC.Data[5596] := 334.81;
   Prof_FEC.Data[5597] := 399.22;
   Prof_FEC.Data[5598] := 395.74;
   Prof_FEC.Data[5599] := 402.22;
   Prof_FEC.Data[5600] := 447.16;
   Prof_FEC.Data[5601] := 516.24;
   Prof_FEC.Data[5602] := 591.52;
   Prof_FEC.Data[5603] := 568.49;
   Prof_FEC.Data[5604] := 626.29;
   Prof_FEC.Data[5605] := 616.52;
   Prof_FEC.Data[5606] := 710.96;
   Prof_FEC.Data[5607] := 701.67;
   Prof_FEC.Data[5608] := 730.81;
   Prof_FEC.Data[5609] := 685.84;
   Prof_FEC.Data[5610] := 730.67;
   Prof_FEC.Data[5611] := 717.44;
   Prof_FEC.Data[5612] := 711.09;
   Prof_FEC.Data[5613] := 705.26;
   Prof_FEC.Data[5614] := 670.48;
   Prof_FEC.Data[5615] := 701.89;
   Prof_FEC.Data[5616] := 595.89;
   Prof_FEC.Data[5617] := 648.8;
   Prof_FEC.Data[5618] := 638.27;
   Prof_FEC.Data[5619] := 581.64;
   Prof_FEC.Data[5620] := 633.38;
   Prof_FEC.Data[5621] := 661.09;
   Prof_FEC.Data[5622] := 641.44;
   Prof_FEC.Data[5623] := 641.46;
   Prof_FEC.Data[5624] := 705.14;
   Prof_FEC.Data[5625] := 614.61;
   Prof_FEC.Data[5626] := 617.56;
   Prof_FEC.Data[5627] := 656.72;
   Prof_FEC.Data[5628] := 720.64;
   Prof_FEC.Data[5629] := 723.6;
   Prof_FEC.Data[5630] := 779.49;
   Prof_FEC.Data[5631] := 803.05;
   Prof_FEC.Data[5632] := 844.1;
   Prof_FEC.Data[5633] := 787.16;
   Prof_FEC.Data[5634] := 703.43;
   Prof_FEC.Data[5635] := 596.31;
   Prof_FEC.Data[5636] := 401.33;
   Prof_FEC.Data[5637] := 321.05;
   Prof_FEC.Data[5638] := 259.2;
   Prof_FEC.Data[5639] := 238.39;
   Prof_FEC.Data[5640] := 257.01;
   Prof_FEC.Data[5641] := 278.45;
   Prof_FEC.Data[5642] := 226.98;
   Prof_FEC.Data[5643] := 242.69;
   Prof_FEC.Data[5644] := 42.363;
   Prof_FEC.Data[5645] := 42.248;
   Prof_FEC.Data[5646] := 41.469;
   Prof_FEC.Data[5647] := 43.164;
   Prof_FEC.Data[5648] := 38.585;
   Prof_FEC.Data[5649] := 41.407;
   Prof_FEC.Data[5650] := 38.687;
   Prof_FEC.Data[5651] := 37.073;
   Prof_FEC.Data[5652] := 37.438;
   Prof_FEC.Data[5653] := 37.608;
   Prof_FEC.Data[5654] := 39.691;
   Prof_FEC.Data[5655] := 42.481;
   Prof_FEC.Data[5656] := 38.911;
   Prof_FEC.Data[5657] := 39.096;
   Prof_FEC.Data[5658] := 38.669;
   Prof_FEC.Data[5659] := 39.993;
   Prof_FEC.Data[5660] := 38.072;
   Prof_FEC.Data[5661] := 40.602;
   Prof_FEC.Data[5662] := 38.051;
   Prof_FEC.Data[5663] := 38.984;
   Prof_FEC.Data[5664] := 37.562;
   Prof_FEC.Data[5665] := 37.603;
   Prof_FEC.Data[5666] := 37.744;
   Prof_FEC.Data[5667] := 35.638;
   Prof_FEC.Data[5668] := 39.976;
   Prof_FEC.Data[5669] := 39.837;
   Prof_FEC.Data[5670] := 38.99;
   Prof_FEC.Data[5671] := 37.41;
   Prof_FEC.Data[5672] := 38.182;
   Prof_FEC.Data[5673] := 38.93;
   Prof_FEC.Data[5674] := 39.306;
   Prof_FEC.Data[5675] := 37.579;
   Prof_FEC.Data[5676] := 41.014;
   Prof_FEC.Data[5677] := 42.153;
   Prof_FEC.Data[5678] := 40.993;
   Prof_FEC.Data[5679] := 42.808;
   Prof_FEC.Data[5680] := 40.432;
   Prof_FEC.Data[5681] := 40.716;
   Prof_FEC.Data[5682] := 40.309;
   Prof_FEC.Data[5683] := 39.813;
   Prof_FEC.Data[5684] := 256.54;
   Prof_FEC.Data[5685] := 242.32;
   Prof_FEC.Data[5686] := 285.55;
   Prof_FEC.Data[5687] := 290.61;
   Prof_FEC.Data[5688] := 282.03;
   Prof_FEC.Data[5689] := 264.46;
   Prof_FEC.Data[5690] := 288.2;
   Prof_FEC.Data[5691] := 285.84;
   Prof_FEC.Data[5692] := 306.36;
   Prof_FEC.Data[5693] := 325.09;
   Prof_FEC.Data[5694] := 327.09;
   Prof_FEC.Data[5695] := 321.55;
   Prof_FEC.Data[5696] := 317.12;
   Prof_FEC.Data[5697] := 310.99;
   Prof_FEC.Data[5698] := 314.57;
   Prof_FEC.Data[5699] := 368.32;
   Prof_FEC.Data[5700] := 389.09;
   Prof_FEC.Data[5701] := 420.38;
   Prof_FEC.Data[5702] := 402.73;
   Prof_FEC.Data[5703] := 405.11;
   Prof_FEC.Data[5704] := 377.69;
   Prof_FEC.Data[5705] := 363.81;
   Prof_FEC.Data[5706] := 418.05;
   Prof_FEC.Data[5707] := 332.91;
   Prof_FEC.Data[5708] := 379.34;
   Prof_FEC.Data[5709] := 400.06;
   Prof_FEC.Data[5710] := 422.72;
   Prof_FEC.Data[5711] := 375.05;
   Prof_FEC.Data[5712] := 355.65;
   Prof_FEC.Data[5713] := 311.73;
   Prof_FEC.Data[5714] := 316.94;
   Prof_FEC.Data[5715] := 314.03;
   Prof_FEC.Data[5716] := 333.11;
   Prof_FEC.Data[5717] := 324.29;
   Prof_FEC.Data[5718] := 335.95;
   Prof_FEC.Data[5719] := 311.9;
   Prof_FEC.Data[5720] := 323.59;
   Prof_FEC.Data[5721] := 329.12;
   Prof_FEC.Data[5722] := 296.06;
   Prof_FEC.Data[5723] := 329.88;
   Prof_FEC.Data[5724] := 370.85;
   Prof_FEC.Data[5725] := 334.41;
   Prof_FEC.Data[5726] := 311.07;
   Prof_FEC.Data[5727] := 266.27;
   Prof_FEC.Data[5728] := 157.77;
   Prof_FEC.Data[5729] := 104.95;
   Prof_FEC.Data[5730] := 90.61;
   Prof_FEC.Data[5731] := 100.68;
   Prof_FEC.Data[5732] := 136.31;
   Prof_FEC.Data[5733] := 133.53;
   Prof_FEC.Data[5734] := 147.34;
   Prof_FEC.Data[5735] := 186.08;
   Prof_FEC.Data[5736] := 217.41;
   Prof_FEC.Data[5737] := 241.95;
   Prof_FEC.Data[5738] := 260.24;
   Prof_FEC.Data[5739] := 279.85;
   Prof_FEC.Data[5740] := 36.508;
   Prof_FEC.Data[5741] := 36.709;
   Prof_FEC.Data[5742] := 37.851;
   Prof_FEC.Data[5743] := 38.309;
   Prof_FEC.Data[5744] := 38.399;
   Prof_FEC.Data[5745] := 38.527;
   Prof_FEC.Data[5746] := 40.289;
   Prof_FEC.Data[5747] := 37.785;
   Prof_FEC.Data[5748] := 38.788;
   Prof_FEC.Data[5749] := 41.268;
   Prof_FEC.Data[5750] := 37.735;
   Prof_FEC.Data[5751] := 39.828;
   Prof_FEC.Data[5752] := 41.218;
   Prof_FEC.Data[5753] := 42.809;
   Prof_FEC.Data[5754] := 45.634;
   Prof_FEC.Data[5755] := 41.892;
   Prof_FEC.Data[5756] := 40.157;
   Prof_FEC.Data[5757] := 41.163;
   Prof_FEC.Data[5758] := 39.465;
   Prof_FEC.Data[5759] := 41.831;
   Prof_FEC.Data[5760] := 41.639;
   Prof_FEC.Data[5761] := 42.334;
   Prof_FEC.Data[5762] := 39.6;
   Prof_FEC.Data[5763] := 42.16;
   Prof_FEC.Data[5764] := 41.401;
   Prof_FEC.Data[5765] := 39.822;
   Prof_FEC.Data[5766] := 38.153;
   Prof_FEC.Data[5767] := 40.271;
   Prof_FEC.Data[5768] := 42.995;
   Prof_FEC.Data[5769] := 42.586;
   Prof_FEC.Data[5770] := 41.465;
   Prof_FEC.Data[5771] := 42.316;
   Prof_FEC.Data[5772] := 41.437;
   Prof_FEC.Data[5773] := 40.015;
   Prof_FEC.Data[5774] := 40.398;
   Prof_FEC.Data[5775] := 39.23;
   Prof_FEC.Data[5776] := 39.5;
   Prof_FEC.Data[5777] := 37.81;
   Prof_FEC.Data[5778] := 39.655;
   Prof_FEC.Data[5779] := 41.463;
   Prof_FEC.Data[5780] := 240.54;
   Prof_FEC.Data[5781] := 238.44;
   Prof_FEC.Data[5782] := 224.87;
   Prof_FEC.Data[5783] := 248.09;
   Prof_FEC.Data[5784] := 260.25;
   Prof_FEC.Data[5785] := 277.07;
   Prof_FEC.Data[5786] := 282.7;
   Prof_FEC.Data[5787] := 214.17;
   Prof_FEC.Data[5788] := 146.03;
   Prof_FEC.Data[5789] := 129.02;
   Prof_FEC.Data[5790] := 106.34;
   Prof_FEC.Data[5791] := 114.58;
   Prof_FEC.Data[5792] := 144.85;
   Prof_FEC.Data[5793] := 135.63;
   Prof_FEC.Data[5794] := 157.61;
   Prof_FEC.Data[5795] := 148.3;
   Prof_FEC.Data[5796] := 131.83;
   Prof_FEC.Data[5797] := 144.39;
   Prof_FEC.Data[5798] := 128.35;
   Prof_FEC.Data[5799] := 138.84;
   Prof_FEC.Data[5800] := 161.65;
   Prof_FEC.Data[5801] := 157.79;
   Prof_FEC.Data[5802] := 155.82;
   Prof_FEC.Data[5803] := 146.27;
   Prof_FEC.Data[5804] := 132.3;
   Prof_FEC.Data[5805] := 126.87;
   Prof_FEC.Data[5806] := 131.47;
   Prof_FEC.Data[5807] := 128.49;
   Prof_FEC.Data[5808] := 157.13;
   Prof_FEC.Data[5809] := 163.48;
   Prof_FEC.Data[5810] := 152.81;
   Prof_FEC.Data[5811] := 148.69;
   Prof_FEC.Data[5812] := 129.53;
   Prof_FEC.Data[5813] := 120.54;
   Prof_FEC.Data[5814] := 133.88;
   Prof_FEC.Data[5815] := 141.46;
   Prof_FEC.Data[5816] := 148.86;
   Prof_FEC.Data[5817] := 164.18;
   Prof_FEC.Data[5818] := 147.99;
   Prof_FEC.Data[5819] := 147.12;
   Prof_FEC.Data[5820] := 135.03;
   Prof_FEC.Data[5821] := 124.56;
   Prof_FEC.Data[5822] := 130.06;
   Prof_FEC.Data[5823] := 137.12;
   Prof_FEC.Data[5824] := 129.64;
   Prof_FEC.Data[5825] := 142.14;
   Prof_FEC.Data[5826] := 141.09;
   Prof_FEC.Data[5827] := 142.58;
   Prof_FEC.Data[5828] := 151.11;
   Prof_FEC.Data[5829] := 168.47;
   Prof_FEC.Data[5830] := 156.64;
   Prof_FEC.Data[5831] := 168.36;
   Prof_FEC.Data[5832] := 229.07;
   Prof_FEC.Data[5833] := 283.24;
   Prof_FEC.Data[5834] := 275.46;
   Prof_FEC.Data[5835] := 244.89;
   Prof_FEC.Data[5836] := 39.845;
   Prof_FEC.Data[5837] := 40.505;
   Prof_FEC.Data[5838] := 40.803;
   Prof_FEC.Data[5839] := 40.395;
   Prof_FEC.Data[5840] := 41.993;
   Prof_FEC.Data[5841] := 44.226;
   Prof_FEC.Data[5842] := 42.555;
   Prof_FEC.Data[5843] := 43.754;
   Prof_FEC.Data[5844] := 41.891;
   Prof_FEC.Data[5845] := 42.635;
   Prof_FEC.Data[5846] := 40.396;
   Prof_FEC.Data[5847] := 40.166;
   Prof_FEC.Data[5848] := 42.842;
   Prof_FEC.Data[5849] := 45.54;
   Prof_FEC.Data[5850] := 45.534;
   Prof_FEC.Data[5851] := 46.944;
   Prof_FEC.Data[5852] := 45.058;
   Prof_FEC.Data[5853] := 43.982;
   Prof_FEC.Data[5854] := 42.865;
   Prof_FEC.Data[5855] := 42.728;
   Prof_FEC.Data[5856] := 44.103;
   Prof_FEC.Data[5857] := 48.436;
   Prof_FEC.Data[5858] := 46.443;
   Prof_FEC.Data[5859] := 42.773;
   Prof_FEC.Data[5860] := 44.184;
   Prof_FEC.Data[5861] := 42.644;
   Prof_FEC.Data[5862] := 44.582;
   Prof_FEC.Data[5863] := 42.769;
   Prof_FEC.Data[5864] := 44.625;
   Prof_FEC.Data[5865] := 46.647;
   Prof_FEC.Data[5866] := 46.827;
   Prof_FEC.Data[5867] := 46.272;
   Prof_FEC.Data[5868] := 46.955;
   Prof_FEC.Data[5869] := 46.285;
   Prof_FEC.Data[5870] := 47.26;
   Prof_FEC.Data[5871] := 44.928;
   Prof_FEC.Data[5872] := 45.842;
   Prof_FEC.Data[5873] := 49.501;
   Prof_FEC.Data[5874] := 44.075;
   Prof_FEC.Data[5875] := 44.323;
   Prof_FEC.Data[5876] := 265.97;
   Prof_FEC.Data[5877] := 247.71;
   Prof_FEC.Data[5878] := 270.3;
   Prof_FEC.Data[5879] := 304.23;
   Prof_FEC.Data[5880] := 328.17;
   Prof_FEC.Data[5881] := 387.67;
   Prof_FEC.Data[5882] := 410.88;
   Prof_FEC.Data[5883] := 398.45;
   Prof_FEC.Data[5884] := 375.25;
   Prof_FEC.Data[5885] := 373.93;
   Prof_FEC.Data[5886] := 431.65;
   Prof_FEC.Data[5887] := 390.93;
   Prof_FEC.Data[5888] := 503.08;
   Prof_FEC.Data[5889] := 433.2;
   Prof_FEC.Data[5890] := 478.68;
   Prof_FEC.Data[5891] := 489.05;
   Prof_FEC.Data[5892] := 567.04;
   Prof_FEC.Data[5893] := 573.32;
   Prof_FEC.Data[5894] := 639.7;
   Prof_FEC.Data[5895] := 590.85;
   Prof_FEC.Data[5896] := 564.15;
   Prof_FEC.Data[5897] := 549.64;
   Prof_FEC.Data[5898] := 626.33;
   Prof_FEC.Data[5899] := 522.44;
   Prof_FEC.Data[5900] := 556.86;
   Prof_FEC.Data[5901] := 578.05;
   Prof_FEC.Data[5902] := 644.73;
   Prof_FEC.Data[5903] := 560.3;
   Prof_FEC.Data[5904] := 642.86;
   Prof_FEC.Data[5905] := 592.65;
   Prof_FEC.Data[5906] := 588.54;
   Prof_FEC.Data[5907] := 619.98;
   Prof_FEC.Data[5908] := 631.5;
   Prof_FEC.Data[5909] := 619.75;
   Prof_FEC.Data[5910] := 636.88;
   Prof_FEC.Data[5911] := 658.1;
   Prof_FEC.Data[5912] := 605.21;
   Prof_FEC.Data[5913] := 600.85;
   Prof_FEC.Data[5914] := 647.48;
   Prof_FEC.Data[5915] := 635.93;
   Prof_FEC.Data[5916] := 570.86;
   Prof_FEC.Data[5917] := 626.21;
   Prof_FEC.Data[5918] := 700.64;
   Prof_FEC.Data[5919] := 621.86;
   Prof_FEC.Data[5920] := 641.53;
   Prof_FEC.Data[5921] := 562.1;
   Prof_FEC.Data[5922] := 569.25;
   Prof_FEC.Data[5923] := 444.72;
   Prof_FEC.Data[5924] := 317.1;
   Prof_FEC.Data[5925] := 242.2;
   Prof_FEC.Data[5926] := 202.87;
   Prof_FEC.Data[5927] := 185.84;
   Prof_FEC.Data[5928] := 234.93;
   Prof_FEC.Data[5929] := 215.87;
   Prof_FEC.Data[5930] := 227.8;
   Prof_FEC.Data[5931] := 244.63;
   Prof_FEC.Data[5932] := 41.657;
   Prof_FEC.Data[5933] := 41.975;
   Prof_FEC.Data[5934] := 43.071;
   Prof_FEC.Data[5935] := 42.324;
   Prof_FEC.Data[5936] := 43.125;
   Prof_FEC.Data[5937] := 37.438;
   Prof_FEC.Data[5938] := 39.464;
   Prof_FEC.Data[5939] := 39.12;
   Prof_FEC.Data[5940] := 43.637;
   Prof_FEC.Data[5941] := 42.185;
   Prof_FEC.Data[5942] := 38.915;
   Prof_FEC.Data[5943] := 40.453;
   Prof_FEC.Data[5944] := 40.204;
   Prof_FEC.Data[5945] := 42.038;
   Prof_FEC.Data[5946] := 40.471;
   Prof_FEC.Data[5947] := 40.948;
   Prof_FEC.Data[5948] := 40.834;
   Prof_FEC.Data[5949] := 41.089;
   Prof_FEC.Data[5950] := 43.293;
   Prof_FEC.Data[5951] := 41.525;
   Prof_FEC.Data[5952] := 41.123;
   Prof_FEC.Data[5953] := 39.614;
   Prof_FEC.Data[5954] := 40.826;
   Prof_FEC.Data[5955] := 38.823;
   Prof_FEC.Data[5956] := 41.929;
   Prof_FEC.Data[5957] := 40.19;
   Prof_FEC.Data[5958] := 43.124;
   Prof_FEC.Data[5959] := 41.74;
   Prof_FEC.Data[5960] := 40.531;
   Prof_FEC.Data[5961] := 40.388;
   Prof_FEC.Data[5962] := 36.429;
   Prof_FEC.Data[5963] := 39.322;
   Prof_FEC.Data[5964] := 42.355;
   Prof_FEC.Data[5965] := 44.53;
   Prof_FEC.Data[5966] := 43.168;
   Prof_FEC.Data[5967] := 38.788;
   Prof_FEC.Data[5968] := 39.588;
   Prof_FEC.Data[5969] := 39.511;
   Prof_FEC.Data[5970] := 40.346;
   Prof_FEC.Data[5971] := 40.057;
   Prof_FEC.Data[5972] := 224.12;
   Prof_FEC.Data[5973] := 246.16;
   Prof_FEC.Data[5974] := 260.0;
   Prof_FEC.Data[5975] := 275.66;
   Prof_FEC.Data[5976] := 366.91;
   Prof_FEC.Data[5977] := 383.03;
   Prof_FEC.Data[5978] := 416.25;
   Prof_FEC.Data[5979] := 427.27;
   Prof_FEC.Data[5980] := 418.12;
   Prof_FEC.Data[5981] := 445.17;
   Prof_FEC.Data[5982] := 413.96;
   Prof_FEC.Data[5983] := 508.63;
   Prof_FEC.Data[5984] := 569.45;
   Prof_FEC.Data[5985] := 612.47;
   Prof_FEC.Data[5986] := 662.06;
   Prof_FEC.Data[5987] := 658.45;
   Prof_FEC.Data[5988] := 653.2;
   Prof_FEC.Data[5989] := 667.78;
   Prof_FEC.Data[5990] := 635.87;
   Prof_FEC.Data[5991] := 651.58;
   Prof_FEC.Data[5992] := 630.96;
   Prof_FEC.Data[5993] := 728.35;
   Prof_FEC.Data[5994] := 661.42;
   Prof_FEC.Data[5995] := 683.02;
   Prof_FEC.Data[5996] := 710.82;
   Prof_FEC.Data[5997] := 730.04;
   Prof_FEC.Data[5998] := 698.07;
   Prof_FEC.Data[5999] := 673.01;
   Prof_FEC.Data[6000] := 650.87;
   Prof_FEC.Data[6001] := 691.16;
   Prof_FEC.Data[6002] := 638.53;
   Prof_FEC.Data[6003] := 665.1;
   Prof_FEC.Data[6004] := 795.45;
   Prof_FEC.Data[6005] := 742.55;
   Prof_FEC.Data[6006] := 784.47;
   Prof_FEC.Data[6007] := 720.56;
   Prof_FEC.Data[6008] := 699.69;
   Prof_FEC.Data[6009] := 675.51;
   Prof_FEC.Data[6010] := 673.63;
   Prof_FEC.Data[6011] := 599.48;
   Prof_FEC.Data[6012] := 660.93;
   Prof_FEC.Data[6013] := 699.63;
   Prof_FEC.Data[6014] := 673.29;
   Prof_FEC.Data[6015] := 662.04;
   Prof_FEC.Data[6016] := 678.55;
   Prof_FEC.Data[6017] := 703.25;
   Prof_FEC.Data[6018] := 625.46;
   Prof_FEC.Data[6019] := 469.01;
   Prof_FEC.Data[6020] := 261.05;
   Prof_FEC.Data[6021] := 211.41;
   Prof_FEC.Data[6022] := 170.56;
   Prof_FEC.Data[6023] := 180.16;
   Prof_FEC.Data[6024] := 209.54;
   Prof_FEC.Data[6025] := 182.11;
   Prof_FEC.Data[6026] := 205.16;
   Prof_FEC.Data[6027] := 202.07;
   Prof_FEC.Data[6028] := 38.303;
   Prof_FEC.Data[6029] := 36.185;
   Prof_FEC.Data[6030] := 34.281;
   Prof_FEC.Data[6031] := 34.47;
   Prof_FEC.Data[6032] := 34.88;
   Prof_FEC.Data[6033] := 33.286;
   Prof_FEC.Data[6034] := 33.703;
   Prof_FEC.Data[6035] := 33.894;
   Prof_FEC.Data[6036] := 35.291;
   Prof_FEC.Data[6037] := 38.143;
   Prof_FEC.Data[6038] := 38.886;
   Prof_FEC.Data[6039] := 36.702;
   Prof_FEC.Data[6040] := 35.463;
   Prof_FEC.Data[6041] := 35.846;
   Prof_FEC.Data[6042] := 35.285;
   Prof_FEC.Data[6043] := 34.883;
   Prof_FEC.Data[6044] := 36.755;
   Prof_FEC.Data[6045] := 38.436;
   Prof_FEC.Data[6046] := 38.416;
   Prof_FEC.Data[6047] := 35.945;
   Prof_FEC.Data[6048] := 37.416;
   Prof_FEC.Data[6049] := 36.795;
   Prof_FEC.Data[6050] := 38.932;
   Prof_FEC.Data[6051] := 37.504;
   Prof_FEC.Data[6052] := 38.477;
   Prof_FEC.Data[6053] := 39.34;
   Prof_FEC.Data[6054] := 40.597;
   Prof_FEC.Data[6055] := 40.868;
   Prof_FEC.Data[6056] := 39.271;
   Prof_FEC.Data[6057] := 39.489;
   Prof_FEC.Data[6058] := 39.565;
   Prof_FEC.Data[6059] := 36.238;
   Prof_FEC.Data[6060] := 39.175;
   Prof_FEC.Data[6061] := 38.955;
   Prof_FEC.Data[6062] := 38.276;
   Prof_FEC.Data[6063] := 39.976;
   Prof_FEC.Data[6064] := 39.768;
   Prof_FEC.Data[6065] := 41.819;
   Prof_FEC.Data[6066] := 38.375;
   Prof_FEC.Data[6067] := 40.692;
   Prof_FEC.Data[6068] := 265.69;
   Prof_FEC.Data[6069] := 257.71;
   Prof_FEC.Data[6070] := 216.42;
   Prof_FEC.Data[6071] := 336.7;
   Prof_FEC.Data[6072] := 372.69;
   Prof_FEC.Data[6073] := 329.78;
   Prof_FEC.Data[6074] := 401.17;
   Prof_FEC.Data[6075] := 449.57;
   Prof_FEC.Data[6076] := 420.51;
   Prof_FEC.Data[6077] := 431.86;
   Prof_FEC.Data[6078] := 476.86;
   Prof_FEC.Data[6079] := 555.03;
   Prof_FEC.Data[6080] := 586.76;
   Prof_FEC.Data[6081] := 625.74;
   Prof_FEC.Data[6082] := 670.56;
   Prof_FEC.Data[6083] := 605.44;
   Prof_FEC.Data[6084] := 600.44;
   Prof_FEC.Data[6085] := 666.81;
   Prof_FEC.Data[6086] := 679.07;
   Prof_FEC.Data[6087] := 685.67;
   Prof_FEC.Data[6088] := 614.53;
   Prof_FEC.Data[6089] := 682.54;
   Prof_FEC.Data[6090] := 722.73;
   Prof_FEC.Data[6091] := 673.46;
   Prof_FEC.Data[6092] := 684.8;
   Prof_FEC.Data[6093] := 680.16;
   Prof_FEC.Data[6094] := 666.31;
   Prof_FEC.Data[6095] := 649.03;
   Prof_FEC.Data[6096] := 571.42;
   Prof_FEC.Data[6097] := 621.75;
   Prof_FEC.Data[6098] := 583.34;
   Prof_FEC.Data[6099] := 644.14;
   Prof_FEC.Data[6100] := 634.89;
   Prof_FEC.Data[6101] := 710.29;
   Prof_FEC.Data[6102] := 684.86;
   Prof_FEC.Data[6103] := 720.53;
   Prof_FEC.Data[6104] := 667.01;
   Prof_FEC.Data[6105] := 661.46;
   Prof_FEC.Data[6106] := 688.85;
   Prof_FEC.Data[6107] := 730.48;
   Prof_FEC.Data[6108] := 682.59;
   Prof_FEC.Data[6109] := 778.26;
   Prof_FEC.Data[6110] := 703.78;
   Prof_FEC.Data[6111] := 664.85;
   Prof_FEC.Data[6112] := 778.14;
   Prof_FEC.Data[6113] := 732.32;
   Prof_FEC.Data[6114] := 677.6;
   Prof_FEC.Data[6115] := 546.22;
   Prof_FEC.Data[6116] := 360.53;
   Prof_FEC.Data[6117] := 289.63;
   Prof_FEC.Data[6118] := 231.85;
   Prof_FEC.Data[6119] := 214.54;
   Prof_FEC.Data[6120] := 252.78;
   Prof_FEC.Data[6121] := 222.1;
   Prof_FEC.Data[6122] := 211.8;
   Prof_FEC.Data[6123] := 232.21;
   Prof_FEC.Data[6124] := 41.07;
   Prof_FEC.Data[6125] := 44.402;
   Prof_FEC.Data[6126] := 41.527;
   Prof_FEC.Data[6127] := 43.272;
   Prof_FEC.Data[6128] := 41.347;
   Prof_FEC.Data[6129] := 44.045;
   Prof_FEC.Data[6130] := 41.632;
   Prof_FEC.Data[6131] := 40.277;
   Prof_FEC.Data[6132] := 42.299;
   Prof_FEC.Data[6133] := 39.856;
   Prof_FEC.Data[6134] := 44.791;
   Prof_FEC.Data[6135] := 40.87;
   Prof_FEC.Data[6136] := 42.911;
   Prof_FEC.Data[6137] := 42.414;
   Prof_FEC.Data[6138] := 41.406;
   Prof_FEC.Data[6139] := 43.405;
   Prof_FEC.Data[6140] := 44.306;
   Prof_FEC.Data[6141] := 43.633;
   Prof_FEC.Data[6142] := 43.273;
   Prof_FEC.Data[6143] := 40.597;
   Prof_FEC.Data[6144] := 40.915;
   Prof_FEC.Data[6145] := 41.474;
   Prof_FEC.Data[6146] := 41.913;
   Prof_FEC.Data[6147] := 43.452;
   Prof_FEC.Data[6148] := 44.641;
   Prof_FEC.Data[6149] := 44.211;
   Prof_FEC.Data[6150] := 45.14;
   Prof_FEC.Data[6151] := 43.167;
   Prof_FEC.Data[6152] := 42.341;
   Prof_FEC.Data[6153] := 43.568;
   Prof_FEC.Data[6154] := 44.854;
   Prof_FEC.Data[6155] := 44.769;
   Prof_FEC.Data[6156] := 47.015;
   Prof_FEC.Data[6157] := 48.87;
   Prof_FEC.Data[6158] := 50.0;
   Prof_FEC.Data[6159] := 49.358;
   Prof_FEC.Data[6160] := 45.871;
   Prof_FEC.Data[6161] := 46.823;
   Prof_FEC.Data[6162] := 49.708;
   Prof_FEC.Data[6163] := 45.881;
   Prof_FEC.Data[6164] := 322.34;
   Prof_FEC.Data[6165] := 309.8;
   Prof_FEC.Data[6166] := 353.9;
   Prof_FEC.Data[6167] := 315.55;
   Prof_FEC.Data[6168] := 358.26;
   Prof_FEC.Data[6169] := 395.46;
   Prof_FEC.Data[6170] := 399.83;
   Prof_FEC.Data[6171] := 397.48;
   Prof_FEC.Data[6172] := 422.89;
   Prof_FEC.Data[6173] := 456.04;
   Prof_FEC.Data[6174] := 467.06;
   Prof_FEC.Data[6175] := 547.14;
   Prof_FEC.Data[6176] := 502.07;
   Prof_FEC.Data[6177] := 580.94;
   Prof_FEC.Data[6178] := 600.03;
   Prof_FEC.Data[6179] := 651.08;
   Prof_FEC.Data[6180] := 703.43;
   Prof_FEC.Data[6181] := 732.29;
   Prof_FEC.Data[6182] := 743.98;
   Prof_FEC.Data[6183] := 780.18;
   Prof_FEC.Data[6184] := 731.71;
   Prof_FEC.Data[6185] := 674.61;
   Prof_FEC.Data[6186] := 683.31;
   Prof_FEC.Data[6187] := 742.83;
   Prof_FEC.Data[6188] := 764.99;
   Prof_FEC.Data[6189] := 712.68;
   Prof_FEC.Data[6190] := 647.19;
   Prof_FEC.Data[6191] := 656.19;
   Prof_FEC.Data[6192] := 625.22;
   Prof_FEC.Data[6193] := 560.75;
   Prof_FEC.Data[6194] := 641.68;
   Prof_FEC.Data[6195] := 643.45;
   Prof_FEC.Data[6196] := 713.06;
   Prof_FEC.Data[6197] := 671.5;
   Prof_FEC.Data[6198] := 664.46;
   Prof_FEC.Data[6199] := 695.84;
   Prof_FEC.Data[6200] := 705.28;
   Prof_FEC.Data[6201] := 636.01;
   Prof_FEC.Data[6202] := 681.15;
   Prof_FEC.Data[6203] := 746.81;
   Prof_FEC.Data[6204] := 710.47;
   Prof_FEC.Data[6205] := 667.24;
   Prof_FEC.Data[6206] := 630.58;
   Prof_FEC.Data[6207] := 701.46;
   Prof_FEC.Data[6208] := 653.53;
   Prof_FEC.Data[6209] := 685.96;
   Prof_FEC.Data[6210] := 669.56;
   Prof_FEC.Data[6211] := 605.69;
   Prof_FEC.Data[6212] := 420.16;
   Prof_FEC.Data[6213] := 309.17;
   Prof_FEC.Data[6214] := 250.53;
   Prof_FEC.Data[6215] := 240.48;
   Prof_FEC.Data[6216] := 269.21;
   Prof_FEC.Data[6217] := 247.0;
   Prof_FEC.Data[6218] := 251.35;
   Prof_FEC.Data[6219] := 236.46;
   Prof_FEC.Data[6220] := 41.7;
   Prof_FEC.Data[6221] := 41.282;
   Prof_FEC.Data[6222] := 42.496;
   Prof_FEC.Data[6223] := 40.912;
   Prof_FEC.Data[6224] := 42.027;
   Prof_FEC.Data[6225] := 40.564;
   Prof_FEC.Data[6226] := 39.572;
   Prof_FEC.Data[6227] := 40.655;
   Prof_FEC.Data[6228] := 45.97;
   Prof_FEC.Data[6229] := 49.788;
   Prof_FEC.Data[6230] := 49.116;
   Prof_FEC.Data[6231] := 45.864;
   Prof_FEC.Data[6232] := 47.644;
   Prof_FEC.Data[6233] := 46.916;
   Prof_FEC.Data[6234] := 49.193;
   Prof_FEC.Data[6235] := 47.291;
   Prof_FEC.Data[6236] := 50.0;
   Prof_FEC.Data[6237] := 49.973;
   Prof_FEC.Data[6238] := 47.131;
   Prof_FEC.Data[6239] := 45.97;
   Prof_FEC.Data[6240] := 46.271;
   Prof_FEC.Data[6241] := 42.81;
   Prof_FEC.Data[6242] := 44.138;
   Prof_FEC.Data[6243] := 49.096;
   Prof_FEC.Data[6244] := 50.0;
   Prof_FEC.Data[6245] := 50.0;
   Prof_FEC.Data[6246] := 50.0;
   Prof_FEC.Data[6247] := 50.0;
   Prof_FEC.Data[6248] := 50.0;
   Prof_FEC.Data[6249] := 45.154;
   Prof_FEC.Data[6250] := 45.087;
   Prof_FEC.Data[6251] := 47.621;
   Prof_FEC.Data[6252] := 50.0;
   Prof_FEC.Data[6253] := 50.0;
   Prof_FEC.Data[6254] := 50.0;
   Prof_FEC.Data[6255] := 50.0;
   Prof_FEC.Data[6256] := 50.0;
   Prof_FEC.Data[6257] := 50.0;
   Prof_FEC.Data[6258] := 48.533;
   Prof_FEC.Data[6259] := 50.0;
   Prof_FEC.Data[6260] := 343.98;
   Prof_FEC.Data[6261] := 377.96;
   Prof_FEC.Data[6262] := 424.01;
   Prof_FEC.Data[6263] := 401.76;
   Prof_FEC.Data[6264] := 431.57;
   Prof_FEC.Data[6265] := 427.35;
   Prof_FEC.Data[6266] := 434.93;
   Prof_FEC.Data[6267] := 428.01;
   Prof_FEC.Data[6268] := 499.17;
   Prof_FEC.Data[6269] := 496.66;
   Prof_FEC.Data[6270] := 500.16;
   Prof_FEC.Data[6271] := 559.3;
   Prof_FEC.Data[6272] := 651.15;
   Prof_FEC.Data[6273] := 617.67;
   Prof_FEC.Data[6274] := 749.72;
   Prof_FEC.Data[6275] := 750.46;
   Prof_FEC.Data[6276] := 834.28;
   Prof_FEC.Data[6277] := 872.39;
   Prof_FEC.Data[6278] := 888.18;
   Prof_FEC.Data[6279] := 852.8;
   Prof_FEC.Data[6280] := 846.21;
   Prof_FEC.Data[6281] := 876.57;
   Prof_FEC.Data[6282] := 826.3;
   Prof_FEC.Data[6283] := 902.77;
   Prof_FEC.Data[6284] := 838.22;
   Prof_FEC.Data[6285] := 805.7;
   Prof_FEC.Data[6286] := 757.08;
   Prof_FEC.Data[6287] := 756.62;
   Prof_FEC.Data[6288] := 765.16;
   Prof_FEC.Data[6289] := 726.33;
   Prof_FEC.Data[6290] := 770.15;
   Prof_FEC.Data[6291] := 690.8;
   Prof_FEC.Data[6292] := 765.36;
   Prof_FEC.Data[6293] := 740.24;
   Prof_FEC.Data[6294] := 880.62;
   Prof_FEC.Data[6295] := 761.3;
   Prof_FEC.Data[6296] := 862.75;
   Prof_FEC.Data[6297] := 775.99;
   Prof_FEC.Data[6298] := 708.05;
   Prof_FEC.Data[6299] := 822.38;
   Prof_FEC.Data[6300] := 772.19;
   Prof_FEC.Data[6301] := 748.43;
   Prof_FEC.Data[6302] := 785.21;
   Prof_FEC.Data[6303] := 771.33;
   Prof_FEC.Data[6304] := 811.1;
   Prof_FEC.Data[6305] := 867.74;
   Prof_FEC.Data[6306] := 821.28;
   Prof_FEC.Data[6307] := 668.86;
   Prof_FEC.Data[6308] := 385.17;
   Prof_FEC.Data[6309] := 300.31;
   Prof_FEC.Data[6310] := 235.66;
   Prof_FEC.Data[6311] := 231.34;
   Prof_FEC.Data[6312] := 279.12;
   Prof_FEC.Data[6313] := 274.43;
   Prof_FEC.Data[6314] := 294.01;
   Prof_FEC.Data[6315] := 262.98;
   Prof_FEC.Data[6316] := 46.381;
   Prof_FEC.Data[6317] := 44.618;
   Prof_FEC.Data[6318] := 40.645;
   Prof_FEC.Data[6319] := 40.895;
   Prof_FEC.Data[6320] := 39.666;
   Prof_FEC.Data[6321] := 40.878;
   Prof_FEC.Data[6322] := 40.506;
   Prof_FEC.Data[6323] := 40.318;
   Prof_FEC.Data[6324] := 41.099;
   Prof_FEC.Data[6325] := 39.965;
   Prof_FEC.Data[6326] := 42.935;
   Prof_FEC.Data[6327] := 39.685;
   Prof_FEC.Data[6328] := 40.421;
   Prof_FEC.Data[6329] := 35.645;
   Prof_FEC.Data[6330] := 38.376;
   Prof_FEC.Data[6331] := 42.03;
   Prof_FEC.Data[6332] := 43.507;
   Prof_FEC.Data[6333] := 46.171;
   Prof_FEC.Data[6334] := 43.086;
   Prof_FEC.Data[6335] := 46.388;
   Prof_FEC.Data[6336] := 43.36;
   Prof_FEC.Data[6337] := 39.723;
   Prof_FEC.Data[6338] := 39.921;
   Prof_FEC.Data[6339] := 42.763;
   Prof_FEC.Data[6340] := 44.391;
   Prof_FEC.Data[6341] := 46.339;
   Prof_FEC.Data[6342] := 47.298;
   Prof_FEC.Data[6343] := 43.811;
   Prof_FEC.Data[6344] := 43.128;
   Prof_FEC.Data[6345] := 42.428;
   Prof_FEC.Data[6346] := 44.161;
   Prof_FEC.Data[6347] := 43.086;
   Prof_FEC.Data[6348] := 47.405;
   Prof_FEC.Data[6349] := 49.719;
   Prof_FEC.Data[6350] := 50.0;
   Prof_FEC.Data[6351] := 47.01;
   Prof_FEC.Data[6352] := 45.635;
   Prof_FEC.Data[6353] := 47.716;
   Prof_FEC.Data[6354] := 45.322;
   Prof_FEC.Data[6355] := 48.095;
   Prof_FEC.Data[6356] := 323.75;
   Prof_FEC.Data[6357] := 365.82;
   Prof_FEC.Data[6358] := 370.17;
   Prof_FEC.Data[6359] := 348.5;
   Prof_FEC.Data[6360] := 280.77;
   Prof_FEC.Data[6361] := 270.88;
   Prof_FEC.Data[6362] := 255.97;
   Prof_FEC.Data[6363] := 267.03;
   Prof_FEC.Data[6364] := 272.05;
   Prof_FEC.Data[6365] := 262.72;
   Prof_FEC.Data[6366] := 273.54;
   Prof_FEC.Data[6367] := 285.69;
   Prof_FEC.Data[6368] := 268.45;
   Prof_FEC.Data[6369] := 272.44;
   Prof_FEC.Data[6370] := 281.44;
   Prof_FEC.Data[6371] := 341.17;
   Prof_FEC.Data[6372] := 324.71;
   Prof_FEC.Data[6373] := 372.32;
   Prof_FEC.Data[6374] := 329.5;
   Prof_FEC.Data[6375] := 305.68;
   Prof_FEC.Data[6376] := 346.44;
   Prof_FEC.Data[6377] := 361.63;
   Prof_FEC.Data[6378] := 343.63;
   Prof_FEC.Data[6379] := 322.57;
   Prof_FEC.Data[6380] := 334.26;
   Prof_FEC.Data[6381] := 346.94;
   Prof_FEC.Data[6382] := 366.35;
   Prof_FEC.Data[6383] := 308.17;
   Prof_FEC.Data[6384] := 271.64;
   Prof_FEC.Data[6385] := 269.44;
   Prof_FEC.Data[6386] := 258.93;
   Prof_FEC.Data[6387] := 286.32;
   Prof_FEC.Data[6388] := 259.31;
   Prof_FEC.Data[6389] := 248.92;
   Prof_FEC.Data[6390] := 236.65;
   Prof_FEC.Data[6391] := 234.47;
   Prof_FEC.Data[6392] := 277.02;
   Prof_FEC.Data[6393] := 247.37;
   Prof_FEC.Data[6394] := 249.42;
   Prof_FEC.Data[6395] := 230.01;
   Prof_FEC.Data[6396] := 260.05;
   Prof_FEC.Data[6397] := 276.1;
   Prof_FEC.Data[6398] := 278.27;
   Prof_FEC.Data[6399] := 196.57;
   Prof_FEC.Data[6400] := 143.86;
   Prof_FEC.Data[6401] := 119.35;
   Prof_FEC.Data[6402] := 114.36;
   Prof_FEC.Data[6403] := 110.53;
   Prof_FEC.Data[6404] := 121.11;
   Prof_FEC.Data[6405] := 107.64;
   Prof_FEC.Data[6406] := 118.53;
   Prof_FEC.Data[6407] := 148.59;
   Prof_FEC.Data[6408] := 198.95;
   Prof_FEC.Data[6409] := 249.14;
   Prof_FEC.Data[6410] := 244.75;
   Prof_FEC.Data[6411] := 257.68;
   Prof_FEC.Data[6412] := 38.665;
   Prof_FEC.Data[6413] := 36.441;
   Prof_FEC.Data[6414] := 38.796;
   Prof_FEC.Data[6415] := 38.581;
   Prof_FEC.Data[6416] := 44.682;
   Prof_FEC.Data[6417] := 44.906;
   Prof_FEC.Data[6418] := 42.205;
   Prof_FEC.Data[6419] := 44.108;
   Prof_FEC.Data[6420] := 39.276;
   Prof_FEC.Data[6421] := 42.252;
   Prof_FEC.Data[6422] := 40.496;
   Prof_FEC.Data[6423] := 39.313;
   Prof_FEC.Data[6424] := 43.082;
   Prof_FEC.Data[6425] := 44.727;
   Prof_FEC.Data[6426] := 45.234;
   Prof_FEC.Data[6427] := 42.094;
   Prof_FEC.Data[6428] := 41.114;
   Prof_FEC.Data[6429] := 40.866;
   Prof_FEC.Data[6430] := 39.112;
   Prof_FEC.Data[6431] := 42.892;
   Prof_FEC.Data[6432] := 46.339;
   Prof_FEC.Data[6433] := 46.144;
   Prof_FEC.Data[6434] := 43.817;
   Prof_FEC.Data[6435] := 42.305;
   Prof_FEC.Data[6436] := 39.43;
   Prof_FEC.Data[6437] := 40.606;
   Prof_FEC.Data[6438] := 44.964;
   Prof_FEC.Data[6439] := 43.199;
   Prof_FEC.Data[6440] := 46.154;
   Prof_FEC.Data[6441] := 45.891;
   Prof_FEC.Data[6442] := 44.776;
   Prof_FEC.Data[6443] := 43.701;
   Prof_FEC.Data[6444] := 43.343;
   Prof_FEC.Data[6445] := 39.965;
   Prof_FEC.Data[6446] := 42.444;
   Prof_FEC.Data[6447] := 41.435;
   Prof_FEC.Data[6448] := 45.786;
   Prof_FEC.Data[6449] := 46.782;
   Prof_FEC.Data[6450] := 50.0;
   Prof_FEC.Data[6451] := 44.222;
   Prof_FEC.Data[6452] := 330.83;
   Prof_FEC.Data[6453] := 270.09;
   Prof_FEC.Data[6454] := 265.8;
   Prof_FEC.Data[6455] := 260.31;
   Prof_FEC.Data[6456] := 280.82;
   Prof_FEC.Data[6457] := 289.42;
   Prof_FEC.Data[6458] := 271.58;
   Prof_FEC.Data[6459] := 240.22;
   Prof_FEC.Data[6460] := 183.17;
   Prof_FEC.Data[6461] := 147.22;
   Prof_FEC.Data[6462] := 144.85;
   Prof_FEC.Data[6463] := 142.89;
   Prof_FEC.Data[6464] := 183.19;
   Prof_FEC.Data[6465] := 181.67;
   Prof_FEC.Data[6466] := 177.24;
   Prof_FEC.Data[6467] := 127.06;
   Prof_FEC.Data[6468] := 114.25;
   Prof_FEC.Data[6469] := 120.0;
   Prof_FEC.Data[6470] := 123.01;
   Prof_FEC.Data[6471] := 133.42;
   Prof_FEC.Data[6472] := 170.67;
   Prof_FEC.Data[6473] := 172.32;
   Prof_FEC.Data[6474] := 164.13;
   Prof_FEC.Data[6475] := 136.71;
   Prof_FEC.Data[6476] := 121.69;
   Prof_FEC.Data[6477] := 123.02;
   Prof_FEC.Data[6478] := 126.8;
   Prof_FEC.Data[6479] := 124.42;
   Prof_FEC.Data[6480] := 157.59;
   Prof_FEC.Data[6481] := 138.81;
   Prof_FEC.Data[6482] := 135.88;
   Prof_FEC.Data[6483] := 143.21;
   Prof_FEC.Data[6484] := 140.24;
   Prof_FEC.Data[6485] := 131.95;
   Prof_FEC.Data[6486] := 109.66;
   Prof_FEC.Data[6487] := 121.64;
   Prof_FEC.Data[6488] := 153.68;
   Prof_FEC.Data[6489] := 150.38;
   Prof_FEC.Data[6490] := 162.0;
   Prof_FEC.Data[6491] := 162.37;
   Prof_FEC.Data[6492] := 149.95;
   Prof_FEC.Data[6493] := 129.25;
   Prof_FEC.Data[6494] := 135.14;
   Prof_FEC.Data[6495] := 149.36;
   Prof_FEC.Data[6496] := 151.71;
   Prof_FEC.Data[6497] := 152.33;
   Prof_FEC.Data[6498] := 154.1;
   Prof_FEC.Data[6499] := 151.98;
   Prof_FEC.Data[6500] := 132.28;
   Prof_FEC.Data[6501] := 128.8;
   Prof_FEC.Data[6502] := 134.86;
   Prof_FEC.Data[6503] := 159.58;
   Prof_FEC.Data[6504] := 224.25;
   Prof_FEC.Data[6505] := 286.63;
   Prof_FEC.Data[6506] := 330.22;
   Prof_FEC.Data[6507] := 306.01;
   Prof_FEC.Data[6508] := 42.375;
   Prof_FEC.Data[6509] := 42.021;
   Prof_FEC.Data[6510] := 43.877;
   Prof_FEC.Data[6511] := 45.685;
   Prof_FEC.Data[6512] := 45.916;
   Prof_FEC.Data[6513] := 45.701;
   Prof_FEC.Data[6514] := 45.305;
   Prof_FEC.Data[6515] := 46.12;
   Prof_FEC.Data[6516] := 43.828;
   Prof_FEC.Data[6517] := 41.926;
   Prof_FEC.Data[6518] := 42.59;
   Prof_FEC.Data[6519] := 42.039;
   Prof_FEC.Data[6520] := 40.978;
   Prof_FEC.Data[6521] := 42.072;
   Prof_FEC.Data[6522] := 45.15;
   Prof_FEC.Data[6523] := 45.865;
   Prof_FEC.Data[6524] := 44.687;
   Prof_FEC.Data[6525] := 42.417;
   Prof_FEC.Data[6526] := 43.522;
   Prof_FEC.Data[6527] := 47.08;
   Prof_FEC.Data[6528] := 46.085;
   Prof_FEC.Data[6529] := 47.702;
   Prof_FEC.Data[6530] := 49.416;
   Prof_FEC.Data[6531] := 45.774;
   Prof_FEC.Data[6532] := 41.51;
   Prof_FEC.Data[6533] := 43.927;
   Prof_FEC.Data[6534] := 42.035;
   Prof_FEC.Data[6535] := 42.237;
   Prof_FEC.Data[6536] := 45.142;
   Prof_FEC.Data[6537] := 39.891;
   Prof_FEC.Data[6538] := 45.94;
   Prof_FEC.Data[6539] := 45.523;
   Prof_FEC.Data[6540] := 42.699;
   Prof_FEC.Data[6541] := 42.167;
   Prof_FEC.Data[6542] := 40.285;
   Prof_FEC.Data[6543] := 42.945;
   Prof_FEC.Data[6544] := 45.335;
   Prof_FEC.Data[6545] := 45.117;
   Prof_FEC.Data[6546] := 45.058;
   Prof_FEC.Data[6547] := 43.66;
   Prof_FEC.Data[6548] := 271.45;
   Prof_FEC.Data[6549] := 271.01;
   Prof_FEC.Data[6550] := 270.24;
   Prof_FEC.Data[6551] := 299.03;
   Prof_FEC.Data[6552] := 320.04;
   Prof_FEC.Data[6553] := 361.17;
   Prof_FEC.Data[6554] := 411.61;
   Prof_FEC.Data[6555] := 395.94;
   Prof_FEC.Data[6556] := 425.3;
   Prof_FEC.Data[6557] := 420.7;
   Prof_FEC.Data[6558] := 454.07;
   Prof_FEC.Data[6559] := 512.44;
   Prof_FEC.Data[6560] := 535.23;
   Prof_FEC.Data[6561] := 532.66;
   Prof_FEC.Data[6562] := 571.36;
   Prof_FEC.Data[6563] := 489.02;
   Prof_FEC.Data[6564] := 462.03;
   Prof_FEC.Data[6565] := 638.25;
   Prof_FEC.Data[6566] := 602.71;
   Prof_FEC.Data[6567] := 598.86;
   Prof_FEC.Data[6568] := 649.91;
   Prof_FEC.Data[6569] := 577.78;
   Prof_FEC.Data[6570] := 577.15;
   Prof_FEC.Data[6571] := 622.5;
   Prof_FEC.Data[6572] := 618.55;
   Prof_FEC.Data[6573] := 631.19;
   Prof_FEC.Data[6574] := 640.03;
   Prof_FEC.Data[6575] := 650.36;
   Prof_FEC.Data[6576] := 575.15;
   Prof_FEC.Data[6577] := 557.87;
   Prof_FEC.Data[6578] := 532.74;
   Prof_FEC.Data[6579] := 553.52;
   Prof_FEC.Data[6580] := 684.27;
   Prof_FEC.Data[6581] := 641.33;
   Prof_FEC.Data[6582] := 647.18;
   Prof_FEC.Data[6583] := 596.08;
   Prof_FEC.Data[6584] := 756.02;
   Prof_FEC.Data[6585] := 625.22;
   Prof_FEC.Data[6586] := 618.18;
   Prof_FEC.Data[6587] := 650.81;
   Prof_FEC.Data[6588] := 622.54;
   Prof_FEC.Data[6589] := 630.67;
   Prof_FEC.Data[6590] := 601.14;
   Prof_FEC.Data[6591] := 672.69;
   Prof_FEC.Data[6592] := 744.43;
   Prof_FEC.Data[6593] := 692.94;
   Prof_FEC.Data[6594] := 578.98;
   Prof_FEC.Data[6595] := 531.75;
   Prof_FEC.Data[6596] := 363.35;
   Prof_FEC.Data[6597] := 261.32;
   Prof_FEC.Data[6598] := 226.47;
   Prof_FEC.Data[6599] := 245.12;
   Prof_FEC.Data[6600] := 269.0;
   Prof_FEC.Data[6601] := 260.47;
   Prof_FEC.Data[6602] := 275.85;
   Prof_FEC.Data[6603] := 268.78;
   Prof_FEC.Data[6604] := 45.538;
   Prof_FEC.Data[6605] := 46.728;
   Prof_FEC.Data[6606] := 47.299;
   Prof_FEC.Data[6607] := 46.843;
   Prof_FEC.Data[6608] := 45.97;
   Prof_FEC.Data[6609] := 43.172;
   Prof_FEC.Data[6610] := 41.406;
   Prof_FEC.Data[6611] := 46.063;
   Prof_FEC.Data[6612] := 45.789;
   Prof_FEC.Data[6613] := 45.63;
   Prof_FEC.Data[6614] := 47.856;
   Prof_FEC.Data[6615] := 47.419;
   Prof_FEC.Data[6616] := 42.818;
   Prof_FEC.Data[6617] := 46.229;
   Prof_FEC.Data[6618] := 47.611;
   Prof_FEC.Data[6619] := 46.038;
   Prof_FEC.Data[6620] := 47.319;
   Prof_FEC.Data[6621] := 44.637;
   Prof_FEC.Data[6622] := 49.396;
   Prof_FEC.Data[6623] := 44.381;
   Prof_FEC.Data[6624] := 42.216;
   Prof_FEC.Data[6625] := 43.671;
   Prof_FEC.Data[6626] := 44.587;
   Prof_FEC.Data[6627] := 46.892;
   Prof_FEC.Data[6628] := 47.989;
   Prof_FEC.Data[6629] := 50.0;
   Prof_FEC.Data[6630] := 50.0;
   Prof_FEC.Data[6631] := 50.0;
   Prof_FEC.Data[6632] := 48.621;
   Prof_FEC.Data[6633] := 47.394;
   Prof_FEC.Data[6634] := 47.92;
   Prof_FEC.Data[6635] := 46.014;
   Prof_FEC.Data[6636] := 50.0;
   Prof_FEC.Data[6637] := 50.0;
   Prof_FEC.Data[6638] := 50.0;
   Prof_FEC.Data[6639] := 50.0;
   Prof_FEC.Data[6640] := 47.535;
   Prof_FEC.Data[6641] := 45.604;
   Prof_FEC.Data[6642] := 49.234;
   Prof_FEC.Data[6643] := 47.281;
   Prof_FEC.Data[6644] := 332.41;
   Prof_FEC.Data[6645] := 320.76;
   Prof_FEC.Data[6646] := 318.16;
   Prof_FEC.Data[6647] := 331.05;
   Prof_FEC.Data[6648] := 338.88;
   Prof_FEC.Data[6649] := 306.03;
   Prof_FEC.Data[6650] := 358.68;
   Prof_FEC.Data[6651] := 402.3;
   Prof_FEC.Data[6652] := 351.27;
   Prof_FEC.Data[6653] := 391.96;
   Prof_FEC.Data[6654] := 469.09;
   Prof_FEC.Data[6655] := 454.97;
   Prof_FEC.Data[6656] := 482.89;
   Prof_FEC.Data[6657] := 617.37;
   Prof_FEC.Data[6658] := 603.89;
   Prof_FEC.Data[6659] := 631.46;
   Prof_FEC.Data[6660] := 638.99;
   Prof_FEC.Data[6661] := 728.65;
   Prof_FEC.Data[6662] := 788.31;
   Prof_FEC.Data[6663] := 686.35;
   Prof_FEC.Data[6664] := 721.32;
   Prof_FEC.Data[6665] := 748.0;
   Prof_FEC.Data[6666] := 790.49;
   Prof_FEC.Data[6667] := 708.22;
   Prof_FEC.Data[6668] := 781.97;
   Prof_FEC.Data[6669] := 721.01;
   Prof_FEC.Data[6670] := 722.78;
   Prof_FEC.Data[6671] := 687.08;
   Prof_FEC.Data[6672] := 631.85;
   Prof_FEC.Data[6673] := 599.49;
   Prof_FEC.Data[6674] := 612.16;
   Prof_FEC.Data[6675] := 607.52;
   Prof_FEC.Data[6676] := 655.38;
   Prof_FEC.Data[6677] := 642.43;
   Prof_FEC.Data[6678] := 673.13;
   Prof_FEC.Data[6679] := 635.44;
   Prof_FEC.Data[6680] := 630.08;
   Prof_FEC.Data[6681] := 585.23;
   Prof_FEC.Data[6682] := 594.73;
   Prof_FEC.Data[6683] := 564.32;
   Prof_FEC.Data[6684] := 657.37;
   Prof_FEC.Data[6685] := 680.26;
   Prof_FEC.Data[6686] := 628.83;
   Prof_FEC.Data[6687] := 611.98;
   Prof_FEC.Data[6688] := 684.47;
   Prof_FEC.Data[6689] := 742.13;
   Prof_FEC.Data[6690] := 674.73;
   Prof_FEC.Data[6691] := 590.09;
   Prof_FEC.Data[6692] := 372.24;
   Prof_FEC.Data[6693] := 275.97;
   Prof_FEC.Data[6694] := 229.71;
   Prof_FEC.Data[6695] := 238.09;
   Prof_FEC.Data[6696] := 269.14;
   Prof_FEC.Data[6697] := 267.07;
   Prof_FEC.Data[6698] := 290.0;
   Prof_FEC.Data[6699] := 320.23;
   Prof_FEC.Data[6700] := 48.338;
   Prof_FEC.Data[6701] := 47.968;
   Prof_FEC.Data[6702] := 47.574;
   Prof_FEC.Data[6703] := 46.062;
   Prof_FEC.Data[6704] := 44.996;
   Prof_FEC.Data[6705] := 42.465;
   Prof_FEC.Data[6706] := 41.558;
   Prof_FEC.Data[6707] := 43.902;
   Prof_FEC.Data[6708] := 46.322;
   Prof_FEC.Data[6709] := 47.375;
   Prof_FEC.Data[6710] := 49.235;
   Prof_FEC.Data[6711] := 47.883;
   Prof_FEC.Data[6712] := 48.156;
   Prof_FEC.Data[6713] := 44.48;
   Prof_FEC.Data[6714] := 45.705;
   Prof_FEC.Data[6715] := 45.566;
   Prof_FEC.Data[6716] := 48.869;
   Prof_FEC.Data[6717] := 47.007;
   Prof_FEC.Data[6718] := 46.865;
   Prof_FEC.Data[6719] := 42.446;
   Prof_FEC.Data[6720] := 42.266;
   Prof_FEC.Data[6721] := 39.673;
   Prof_FEC.Data[6722] := 38.78;
   Prof_FEC.Data[6723] := 42.769;
   Prof_FEC.Data[6724] := 41.199;
   Prof_FEC.Data[6725] := 43.453;
   Prof_FEC.Data[6726] := 44.208;
   Prof_FEC.Data[6727] := 43.128;
   Prof_FEC.Data[6728] := 40.64;
   Prof_FEC.Data[6729] := 41.2;
   Prof_FEC.Data[6730] := 42.023;
   Prof_FEC.Data[6731] := 41.916;
   Prof_FEC.Data[6732] := 48.478;
   Prof_FEC.Data[6733] := 44.92;
   Prof_FEC.Data[6734] := 43.999;
   Prof_FEC.Data[6735] := 42.324;
   Prof_FEC.Data[6736] := 45.052;
   Prof_FEC.Data[6737] := 40.82;
   Prof_FEC.Data[6738] := 42.538;
   Prof_FEC.Data[6739] := 42.681;
   Prof_FEC.Data[6740] := 315.73;
   Prof_FEC.Data[6741] := 340.79;
   Prof_FEC.Data[6742] := 327.55;
   Prof_FEC.Data[6743] := 354.29;
   Prof_FEC.Data[6744] := 332.79;
   Prof_FEC.Data[6745] := 398.82;
   Prof_FEC.Data[6746] := 434.6;
   Prof_FEC.Data[6747] := 433.5;
   Prof_FEC.Data[6748] := 460.84;
   Prof_FEC.Data[6749] := 405.59;
   Prof_FEC.Data[6750] := 484.67;
   Prof_FEC.Data[6751] := 530.69;
   Prof_FEC.Data[6752] := 568.18;
   Prof_FEC.Data[6753] := 634.7;
   Prof_FEC.Data[6754] := 664.21;
   Prof_FEC.Data[6755] := 681.5;
   Prof_FEC.Data[6756] := 700.95;
   Prof_FEC.Data[6757] := 820.91;
   Prof_FEC.Data[6758] := 693.71;
   Prof_FEC.Data[6759] := 686.04;
   Prof_FEC.Data[6760] := 702.39;
   Prof_FEC.Data[6761] := 657.52;
   Prof_FEC.Data[6762] := 755.02;
   Prof_FEC.Data[6763] := 781.66;
   Prof_FEC.Data[6764] := 679.15;
   Prof_FEC.Data[6765] := 676.86;
   Prof_FEC.Data[6766] := 615.41;
   Prof_FEC.Data[6767] := 671.35;
   Prof_FEC.Data[6768] := 550.59;
   Prof_FEC.Data[6769] := 606.49;
   Prof_FEC.Data[6770] := 675.29;
   Prof_FEC.Data[6771] := 666.8;
   Prof_FEC.Data[6772] := 619.28;
   Prof_FEC.Data[6773] := 668.44;
   Prof_FEC.Data[6774] := 633.54;
   Prof_FEC.Data[6775] := 646.97;
   Prof_FEC.Data[6776] := 633.67;
   Prof_FEC.Data[6777] := 638.65;
   Prof_FEC.Data[6778] := 720.14;
   Prof_FEC.Data[6779] := 699.44;
   Prof_FEC.Data[6780] := 730.03;
   Prof_FEC.Data[6781] := 676.89;
   Prof_FEC.Data[6782] := 681.58;
   Prof_FEC.Data[6783] := 671.65;
   Prof_FEC.Data[6784] := 731.22;
   Prof_FEC.Data[6785] := 744.4;
   Prof_FEC.Data[6786] := 656.64;
   Prof_FEC.Data[6787] := 530.7;
   Prof_FEC.Data[6788] := 364.66;
   Prof_FEC.Data[6789] := 287.02;
   Prof_FEC.Data[6790] := 224.9;
   Prof_FEC.Data[6791] := 234.55;
   Prof_FEC.Data[6792] := 229.81;
   Prof_FEC.Data[6793] := 236.09;
   Prof_FEC.Data[6794] := 248.28;
   Prof_FEC.Data[6795] := 266.59;
   Prof_FEC.Data[6796] := 44.027;
   Prof_FEC.Data[6797] := 44.362;
   Prof_FEC.Data[6798] := 42.936;
   Prof_FEC.Data[6799] := 41.321;
   Prof_FEC.Data[6800] := 40.625;
   Prof_FEC.Data[6801] := 41.899;
   Prof_FEC.Data[6802] := 40.116;
   Prof_FEC.Data[6803] := 41.914;
   Prof_FEC.Data[6804] := 45.524;
   Prof_FEC.Data[6805] := 48.601;
   Prof_FEC.Data[6806] := 43.363;
   Prof_FEC.Data[6807] := 43.237;
   Prof_FEC.Data[6808] := 40.022;
   Prof_FEC.Data[6809] := 41.811;
   Prof_FEC.Data[6810] := 44.341;
   Prof_FEC.Data[6811] := 45.3;
   Prof_FEC.Data[6812] := 46.039;
   Prof_FEC.Data[6813] := 45.757;
   Prof_FEC.Data[6814] := 46.241;
   Prof_FEC.Data[6815] := 43.314;
   Prof_FEC.Data[6816] := 45.185;
   Prof_FEC.Data[6817] := 42.537;
   Prof_FEC.Data[6818] := 44.946;
   Prof_FEC.Data[6819] := 45.893;
   Prof_FEC.Data[6820] := 49.654;
   Prof_FEC.Data[6821] := 50.0;
   Prof_FEC.Data[6822] := 50.0;
   Prof_FEC.Data[6823] := 50.0;
   Prof_FEC.Data[6824] := 50.0;
   Prof_FEC.Data[6825] := 50.0;
   Prof_FEC.Data[6826] := 47.474;
   Prof_FEC.Data[6827] := 46.861;
   Prof_FEC.Data[6828] := 49.519;
   Prof_FEC.Data[6829] := 50.0;
   Prof_FEC.Data[6830] := 50.0;
   Prof_FEC.Data[6831] := 50.0;
   Prof_FEC.Data[6832] := 49.674;
   Prof_FEC.Data[6833] := 50.0;
   Prof_FEC.Data[6834] := 50.0;
   Prof_FEC.Data[6835] := 50.0;
   Prof_FEC.Data[6836] := 376.72;
   Prof_FEC.Data[6837] := 429.55;
   Prof_FEC.Data[6838] := 407.69;
   Prof_FEC.Data[6839] := 390.77;
   Prof_FEC.Data[6840] := 373.33;
   Prof_FEC.Data[6841] := 367.77;
   Prof_FEC.Data[6842] := 412.86;
   Prof_FEC.Data[6843] := 406.65;
   Prof_FEC.Data[6844] := 456.97;
   Prof_FEC.Data[6845] := 453.11;
   Prof_FEC.Data[6846] := 496.77;
   Prof_FEC.Data[6847] := 543.19;
   Prof_FEC.Data[6848] := 620.26;
   Prof_FEC.Data[6849] := 597.88;
   Prof_FEC.Data[6850] := 660.02;
   Prof_FEC.Data[6851] := 660.54;
   Prof_FEC.Data[6852] := 715.68;
   Prof_FEC.Data[6853] := 758.46;
   Prof_FEC.Data[6854] := 806.44;
   Prof_FEC.Data[6855] := 809.31;
   Prof_FEC.Data[6856] := 779.33;
   Prof_FEC.Data[6857] := 727.38;
   Prof_FEC.Data[6858] := 706.58;
   Prof_FEC.Data[6859] := 678.21;
   Prof_FEC.Data[6860] := 656.92;
   Prof_FEC.Data[6861] := 648.17;
   Prof_FEC.Data[6862] := 689.3;
   Prof_FEC.Data[6863] := 610.8;
   Prof_FEC.Data[6864] := 540.78;
   Prof_FEC.Data[6865] := 609.04;
   Prof_FEC.Data[6866] := 599.35;
   Prof_FEC.Data[6867] := 652.93;
   Prof_FEC.Data[6868] := 650.4;
   Prof_FEC.Data[6869] := 625.89;
   Prof_FEC.Data[6870] := 626.9;
   Prof_FEC.Data[6871] := 694.25;
   Prof_FEC.Data[6872] := 688.02;
   Prof_FEC.Data[6873] := 590.93;
   Prof_FEC.Data[6874] := 562.06;
   Prof_FEC.Data[6875] := 636.58;
   Prof_FEC.Data[6876] := 586.5;
   Prof_FEC.Data[6877] := 595.34;
   Prof_FEC.Data[6878] := 616.25;
   Prof_FEC.Data[6879] := 599.55;
   Prof_FEC.Data[6880] := 610.4;
   Prof_FEC.Data[6881] := 667.94;
   Prof_FEC.Data[6882] := 622.65;
   Prof_FEC.Data[6883] := 503.66;
   Prof_FEC.Data[6884] := 384.65;
   Prof_FEC.Data[6885] := 291.8;
   Prof_FEC.Data[6886] := 254.43;
   Prof_FEC.Data[6887] := 259.53;
   Prof_FEC.Data[6888] := 305.22;
   Prof_FEC.Data[6889] := 303.63;
   Prof_FEC.Data[6890] := 304.64;
   Prof_FEC.Data[6891] := 306.81;
   Prof_FEC.Data[6892] := 44.734;
   Prof_FEC.Data[6893] := 43.022;
   Prof_FEC.Data[6894] := 46.44;
   Prof_FEC.Data[6895] := 45.706;
   Prof_FEC.Data[6896] := 42.948;
   Prof_FEC.Data[6897] := 43.175;
   Prof_FEC.Data[6898] := 39.52;
   Prof_FEC.Data[6899] := 39.748;
   Prof_FEC.Data[6900] := 39.738;
   Prof_FEC.Data[6901] := 41.911;
   Prof_FEC.Data[6902] := 40.282;
   Prof_FEC.Data[6903] := 44.147;
   Prof_FEC.Data[6904] := 40.091;
   Prof_FEC.Data[6905] := 41.813;
   Prof_FEC.Data[6906] := 41.066;
   Prof_FEC.Data[6907] := 44.382;
   Prof_FEC.Data[6908] := 46.37;
   Prof_FEC.Data[6909] := 45.638;
   Prof_FEC.Data[6910] := 47.089;
   Prof_FEC.Data[6911] := 47.868;
   Prof_FEC.Data[6912] := 45.382;
   Prof_FEC.Data[6913] := 41.105;
   Prof_FEC.Data[6914] := 41.989;
   Prof_FEC.Data[6915] := 41.201;
   Prof_FEC.Data[6916] := 45.008;
   Prof_FEC.Data[6917] := 45.55;
   Prof_FEC.Data[6918] := 45.67;
   Prof_FEC.Data[6919] := 43.232;
   Prof_FEC.Data[6920] := 41.284;
   Prof_FEC.Data[6921] := 40.175;
   Prof_FEC.Data[6922] := 40.778;
   Prof_FEC.Data[6923] := 39.372;
   Prof_FEC.Data[6924] := 40.501;
   Prof_FEC.Data[6925] := 44.033;
   Prof_FEC.Data[6926] := 44.865;
   Prof_FEC.Data[6927] := 40.516;
   Prof_FEC.Data[6928] := 41.041;
   Prof_FEC.Data[6929] := 42.755;
   Prof_FEC.Data[6930] := 41.615;
   Prof_FEC.Data[6931] := 43.557;
   Prof_FEC.Data[6932] := 268.68;
   Prof_FEC.Data[6933] := 245.97;
   Prof_FEC.Data[6934] := 273.37;
   Prof_FEC.Data[6935] := 282.27;
   Prof_FEC.Data[6936] := 290.91;
   Prof_FEC.Data[6937] := 297.04;
   Prof_FEC.Data[6938] := 314.86;
   Prof_FEC.Data[6939] := 318.41;
   Prof_FEC.Data[6940] := 381.84;
   Prof_FEC.Data[6941] := 359.84;
   Prof_FEC.Data[6942] := 394.24;
   Prof_FEC.Data[6943] := 461.19;
   Prof_FEC.Data[6944] := 500.61;
   Prof_FEC.Data[6945] := 484.75;
   Prof_FEC.Data[6946] := 486.73;
   Prof_FEC.Data[6947] := 550.85;
   Prof_FEC.Data[6948] := 583.01;
   Prof_FEC.Data[6949] := 653.59;
   Prof_FEC.Data[6950] := 656.77;
   Prof_FEC.Data[6951] := 593.91;
   Prof_FEC.Data[6952] := 590.19;
   Prof_FEC.Data[6953] := 597.73;
   Prof_FEC.Data[6954] := 604.43;
   Prof_FEC.Data[6955] := 592.89;
   Prof_FEC.Data[6956] := 644.66;
   Prof_FEC.Data[6957] := 671.65;
   Prof_FEC.Data[6958] := 668.03;
   Prof_FEC.Data[6959] := 629.6;
   Prof_FEC.Data[6960] := 596.88;
   Prof_FEC.Data[6961] := 543.04;
   Prof_FEC.Data[6962] := 551.15;
   Prof_FEC.Data[6963] := 550.4;
   Prof_FEC.Data[6964] := 581.72;
   Prof_FEC.Data[6965] := 592.49;
   Prof_FEC.Data[6966] := 590.32;
   Prof_FEC.Data[6967] := 575.76;
   Prof_FEC.Data[6968] := 575.84;
   Prof_FEC.Data[6969] := 533.51;
   Prof_FEC.Data[6970] := 608.72;
   Prof_FEC.Data[6971] := 617.29;
   Prof_FEC.Data[6972] := 564.42;
   Prof_FEC.Data[6973] := 691.89;
   Prof_FEC.Data[6974] := 643.81;
   Prof_FEC.Data[6975] := 635.83;
   Prof_FEC.Data[6976] := 814.55;
   Prof_FEC.Data[6977] := 748.51;
   Prof_FEC.Data[6978] := 713.43;
   Prof_FEC.Data[6979] := 552.85;
   Prof_FEC.Data[6980] := 302.34;
   Prof_FEC.Data[6981] := 215.89;
   Prof_FEC.Data[6982] := 183.38;
   Prof_FEC.Data[6983] := 187.75;
   Prof_FEC.Data[6984] := 232.3;
   Prof_FEC.Data[6985] := 210.01;
   Prof_FEC.Data[6986] := 243.95;
   Prof_FEC.Data[6987] := 230.76;
   Prof_FEC.Data[6988] := 41.795;
   Prof_FEC.Data[6989] := 39.596;
   Prof_FEC.Data[6990] := 39.578;
   Prof_FEC.Data[6991] := 39.111;
   Prof_FEC.Data[6992] := 40.254;
   Prof_FEC.Data[6993] := 36.329;
   Prof_FEC.Data[6994] := 37.383;
   Prof_FEC.Data[6995] := 36.735;
   Prof_FEC.Data[6996] := 37.518;
   Prof_FEC.Data[6997] := 37.708;
   Prof_FEC.Data[6998] := 40.349;
   Prof_FEC.Data[6999] := 39.425;
   Prof_FEC.Data[7000] := 38.431;
   Prof_FEC.Data[7001] := 38.705;
   Prof_FEC.Data[7002] := 41.486;
   Prof_FEC.Data[7003] := 37.834;
   Prof_FEC.Data[7004] := 41.483;
   Prof_FEC.Data[7005] := 40.362;
   Prof_FEC.Data[7006] := 41.519;
   Prof_FEC.Data[7007] := 39.783;
   Prof_FEC.Data[7008] := 37.727;
   Prof_FEC.Data[7009] := 39.727;
   Prof_FEC.Data[7010] := 38.295;
   Prof_FEC.Data[7011] := 41.268;
   Prof_FEC.Data[7012] := 39.799;
   Prof_FEC.Data[7013] := 41.795;
   Prof_FEC.Data[7014] := 40.701;
   Prof_FEC.Data[7015] := 39.935;
   Prof_FEC.Data[7016] := 37.931;
   Prof_FEC.Data[7017] := 38.183;
   Prof_FEC.Data[7018] := 38.738;
   Prof_FEC.Data[7019] := 38.001;
   Prof_FEC.Data[7020] := 40.385;
   Prof_FEC.Data[7021] := 40.463;
   Prof_FEC.Data[7022] := 39.524;
   Prof_FEC.Data[7023] := 42.005;
   Prof_FEC.Data[7024] := 40.238;
   Prof_FEC.Data[7025] := 36.915;
   Prof_FEC.Data[7026] := 39.303;
   Prof_FEC.Data[7027] := 37.586;
   Prof_FEC.Data[7028] := 247.26;
   Prof_FEC.Data[7029] := 269.91;
   Prof_FEC.Data[7030] := 260.66;
   Prof_FEC.Data[7031] := 234.08;
   Prof_FEC.Data[7032] := 195.78;
   Prof_FEC.Data[7033] := 164.35;
   Prof_FEC.Data[7034] := 168.64;
   Prof_FEC.Data[7035] := 188.31;
   Prof_FEC.Data[7036] := 242.83;
   Prof_FEC.Data[7037] := 208.49;
   Prof_FEC.Data[7038] := 275.17;
   Prof_FEC.Data[7039] := 265.26;
   Prof_FEC.Data[7040] := 248.75;
   Prof_FEC.Data[7041] := 256.38;
   Prof_FEC.Data[7042] := 270.17;
   Prof_FEC.Data[7043] := 267.18;
   Prof_FEC.Data[7044] := 353.68;
   Prof_FEC.Data[7045] := 388.71;
   Prof_FEC.Data[7046] := 326.17;
   Prof_FEC.Data[7047] := 374.64;
   Prof_FEC.Data[7048] := 355.47;
   Prof_FEC.Data[7049] := 317.22;
   Prof_FEC.Data[7050] := 344.57;
   Prof_FEC.Data[7051] := 363.87;
   Prof_FEC.Data[7052] := 332.45;
   Prof_FEC.Data[7053] := 358.37;
   Prof_FEC.Data[7054] := 330.42;
   Prof_FEC.Data[7055] := 339.2;
   Prof_FEC.Data[7056] := 265.36;
   Prof_FEC.Data[7057] := 262.67;
   Prof_FEC.Data[7058] := 255.42;
   Prof_FEC.Data[7059] := 245.95;
   Prof_FEC.Data[7060] := 253.8;
   Prof_FEC.Data[7061] := 274.24;
   Prof_FEC.Data[7062] := 258.17;
   Prof_FEC.Data[7063] := 300.1;
   Prof_FEC.Data[7064] := 293.03;
   Prof_FEC.Data[7065] := 256.42;
   Prof_FEC.Data[7066] := 264.58;
   Prof_FEC.Data[7067] := 262.77;
   Prof_FEC.Data[7068] := 261.56;
   Prof_FEC.Data[7069] := 268.66;
   Prof_FEC.Data[7070] := 265.4;
   Prof_FEC.Data[7071] := 221.41;
   Prof_FEC.Data[7072] := 143.92;
   Prof_FEC.Data[7073] := 121.33;
   Prof_FEC.Data[7074] := 89.0;
   Prof_FEC.Data[7075] := 91.85;
   Prof_FEC.Data[7076] := 83.73;
   Prof_FEC.Data[7077] := 95.83;
   Prof_FEC.Data[7078] := 96.18;
   Prof_FEC.Data[7079] := 138.72;
   Prof_FEC.Data[7080] := 215.98;
   Prof_FEC.Data[7081] := 222.64;
   Prof_FEC.Data[7082] := 261.89;
   Prof_FEC.Data[7083] := 260.61;
   Prof_FEC.Data[7084] := 37.216;
   Prof_FEC.Data[7085] := 38.619;
   Prof_FEC.Data[7086] := 38.243;
   Prof_FEC.Data[7087] := 40.093;
   Prof_FEC.Data[7088] := 42.074;
   Prof_FEC.Data[7089] := 41.498;
   Prof_FEC.Data[7090] := 39.515;
   Prof_FEC.Data[7091] := 40.808;
   Prof_FEC.Data[7092] := 37.225;
   Prof_FEC.Data[7093] := 39.545;
   Prof_FEC.Data[7094] := 40.532;
   Prof_FEC.Data[7095] := 41.795;
   Prof_FEC.Data[7096] := 44.905;
   Prof_FEC.Data[7097] := 42.809;
   Prof_FEC.Data[7098] := 41.266;
   Prof_FEC.Data[7099] := 39.502;
   Prof_FEC.Data[7100] := 39.795;
   Prof_FEC.Data[7101] := 38.438;
   Prof_FEC.Data[7102] := 36.76;
   Prof_FEC.Data[7103] := 39.076;
   Prof_FEC.Data[7104] := 42.131;
   Prof_FEC.Data[7105] := 40.862;
   Prof_FEC.Data[7106] := 39.671;
   Prof_FEC.Data[7107] := 39.894;
   Prof_FEC.Data[7108] := 37.691;
   Prof_FEC.Data[7109] := 35.453;
   Prof_FEC.Data[7110] := 36.736;
   Prof_FEC.Data[7111] := 39.61;
   Prof_FEC.Data[7112] := 42.119;
   Prof_FEC.Data[7113] := 43.569;
   Prof_FEC.Data[7114] := 40.462;
   Prof_FEC.Data[7115] := 42.521;
   Prof_FEC.Data[7116] := 39.918;
   Prof_FEC.Data[7117] := 37.312;
   Prof_FEC.Data[7118] := 38.4;
   Prof_FEC.Data[7119] := 38.951;
   Prof_FEC.Data[7120] := 42.826;
   Prof_FEC.Data[7121] := 45.038;
   Prof_FEC.Data[7122] := 42.653;
   Prof_FEC.Data[7123] := 42.806;
   Prof_FEC.Data[7124] := 262.16;
   Prof_FEC.Data[7125] := 271.99;
   Prof_FEC.Data[7126] := 225.04;
   Prof_FEC.Data[7127] := 239.6;
   Prof_FEC.Data[7128] := 244.3;
   Prof_FEC.Data[7129] := 215.02;
   Prof_FEC.Data[7130] := 194.1;
   Prof_FEC.Data[7131] := 187.79;
   Prof_FEC.Data[7132] := 142.98;
   Prof_FEC.Data[7133] := 122.98;
   Prof_FEC.Data[7134] := 115.19;
   Prof_FEC.Data[7135] := 132.31;
   Prof_FEC.Data[7136] := 132.99;
   Prof_FEC.Data[7137] := 145.9;
   Prof_FEC.Data[7138] := 143.45;
   Prof_FEC.Data[7139] := 124.55;
   Prof_FEC.Data[7140] := 126.86;
   Prof_FEC.Data[7141] := 111.81;
   Prof_FEC.Data[7142] := 113.9;
   Prof_FEC.Data[7143] := 126.81;
   Prof_FEC.Data[7144] := 134.67;
   Prof_FEC.Data[7145] := 141.12;
   Prof_FEC.Data[7146] := 121.21;
   Prof_FEC.Data[7147] := 137.7;
   Prof_FEC.Data[7148] := 119.31;
   Prof_FEC.Data[7149] := 112.17;
   Prof_FEC.Data[7150] := 111.65;
   Prof_FEC.Data[7151] := 116.75;
   Prof_FEC.Data[7152] := 132.27;
   Prof_FEC.Data[7153] := 123.59;
   Prof_FEC.Data[7154] := 133.23;
   Prof_FEC.Data[7155] := 142.94;
   Prof_FEC.Data[7156] := 113.45;
   Prof_FEC.Data[7157] := 117.7;
   Prof_FEC.Data[7158] := 108.64;
   Prof_FEC.Data[7159] := 115.09;
   Prof_FEC.Data[7160] := 127.41;
   Prof_FEC.Data[7161] := 130.92;
   Prof_FEC.Data[7162] := 126.3;
   Prof_FEC.Data[7163] := 120.09;
   Prof_FEC.Data[7164] := 124.01;
   Prof_FEC.Data[7165] := 113.67;
   Prof_FEC.Data[7166] := 111.61;
   Prof_FEC.Data[7167] := 123.12;
   Prof_FEC.Data[7168] := 114.51;
   Prof_FEC.Data[7169] := 128.35;
   Prof_FEC.Data[7170] := 116.38;
   Prof_FEC.Data[7171] := 117.43;
   Prof_FEC.Data[7172] := 80.93;
   Prof_FEC.Data[7173] := 84.79;
   Prof_FEC.Data[7174] := 89.93;
   Prof_FEC.Data[7175] := 123.91;
   Prof_FEC.Data[7176] := 195.86;
   Prof_FEC.Data[7177] := 221.42;
   Prof_FEC.Data[7178] := 227.4;
   Prof_FEC.Data[7179] := 249.3;
   Prof_FEC.Data[7180] := 38.92;
   Prof_FEC.Data[7181] := 39.487;
   Prof_FEC.Data[7182] := 38.933;
   Prof_FEC.Data[7183] := 38.841;
   Prof_FEC.Data[7184] := 39.198;
   Prof_FEC.Data[7185] := 40.562;
   Prof_FEC.Data[7186] := 42.164;
   Prof_FEC.Data[7187] := 40.581;
   Prof_FEC.Data[7188] := 39.454;
   Prof_FEC.Data[7189] := 38.316;
   Prof_FEC.Data[7190] := 39.13;
   Prof_FEC.Data[7191] := 39.441;
   Prof_FEC.Data[7192] := 39.669;
   Prof_FEC.Data[7193] := 39.767;
   Prof_FEC.Data[7194] := 40.617;
   Prof_FEC.Data[7195] := 39.414;
   Prof_FEC.Data[7196] := 39.548;
   Prof_FEC.Data[7197] := 38.522;
   Prof_FEC.Data[7198] := 38.305;
   Prof_FEC.Data[7199] := 38.998;
   Prof_FEC.Data[7200] := 39.328;
   Prof_FEC.Data[7201] := 35.075;
   Prof_FEC.Data[7202] := 38.727;
   Prof_FEC.Data[7203] := 39.858;
   Prof_FEC.Data[7204] := 37.023;
   Prof_FEC.Data[7205] := 37.976;
   Prof_FEC.Data[7206] := 39.852;
   Prof_FEC.Data[7207] := 39.708;
   Prof_FEC.Data[7208] := 40.701;
   Prof_FEC.Data[7209] := 42.694;
   Prof_FEC.Data[7210] := 41.002;
   Prof_FEC.Data[7211] := 39.491;
   Prof_FEC.Data[7212] := 34.811;
   Prof_FEC.Data[7213] := 35.51;
   Prof_FEC.Data[7214] := 35.272;
   Prof_FEC.Data[7215] := 34.253;
   Prof_FEC.Data[7216] := 36.907;
   Prof_FEC.Data[7217] := 35.427;
   Prof_FEC.Data[7218] := 38.893;
   Prof_FEC.Data[7219] := 42.002;
   Prof_FEC.Data[7220] := 346.29;
   Prof_FEC.Data[7221] := 364.45;
   Prof_FEC.Data[7222] := 382.6;
   Prof_FEC.Data[7223] := 447.91;
   Prof_FEC.Data[7224] := 538.15;
   Prof_FEC.Data[7225] := 518.4;
   Prof_FEC.Data[7226] := 542.42;
   Prof_FEC.Data[7227] := 538.26;
   Prof_FEC.Data[7228] := 541.72;
   Prof_FEC.Data[7229] := 569.87;
   Prof_FEC.Data[7230] := 606.48;
   Prof_FEC.Data[7231] := 534.5;
   Prof_FEC.Data[7232] := 546.97;
   Prof_FEC.Data[7233] := 570.08;
   Prof_FEC.Data[7234] := 575.13;
   Prof_FEC.Data[7235] := 652.02;
   Prof_FEC.Data[7236] := 704.23;
   Prof_FEC.Data[7237] := 640.56;
   Prof_FEC.Data[7238] := 512.35;
   Prof_FEC.Data[7239] := 609.39;
   Prof_FEC.Data[7240] := 648.27;
   Prof_FEC.Data[7241] := 646.26;
   Prof_FEC.Data[7242] := 714.15;
   Prof_FEC.Data[7243] := 678.19;
   Prof_FEC.Data[7244] := 661.53;
   Prof_FEC.Data[7245] := 617.02;
   Prof_FEC.Data[7246] := 624.8;
   Prof_FEC.Data[7247] := 672.39;
   Prof_FEC.Data[7248] := 726.23;
   Prof_FEC.Data[7249] := 709.2;
   Prof_FEC.Data[7250] := 690.91;
   Prof_FEC.Data[7251] := 660.61;
   Prof_FEC.Data[7252] := 681.7;
   Prof_FEC.Data[7253] := 656.98;
   Prof_FEC.Data[7254] := 688.51;
   Prof_FEC.Data[7255] := 717.49;
   Prof_FEC.Data[7256] := 717.67;
   Prof_FEC.Data[7257] := 712.73;
   Prof_FEC.Data[7258] := 683.88;
   Prof_FEC.Data[7259] := 625.65;
   Prof_FEC.Data[7260] := 674.98;
   Prof_FEC.Data[7261] := 645.18;
   Prof_FEC.Data[7262] := 588.8;
   Prof_FEC.Data[7263] := 560.61;
   Prof_FEC.Data[7264] := 274.32;
   Prof_FEC.Data[7265] := 191.1;
   Prof_FEC.Data[7266] := 154.62;
   Prof_FEC.Data[7267] := 127.08;
   Prof_FEC.Data[7268] := 113.45;
   Prof_FEC.Data[7269] := 81.41;
   Prof_FEC.Data[7270] := 87.29;
   Prof_FEC.Data[7271] := 102.75;
   Prof_FEC.Data[7272] := 171.44;
   Prof_FEC.Data[7273] := 223.26;
   Prof_FEC.Data[7274] := 231.75;
   Prof_FEC.Data[7275] := 227.34;
   Prof_FEC.Data[7276] := 34.084;
   Prof_FEC.Data[7277] := 36.6;
   Prof_FEC.Data[7278] := 36.206;
   Prof_FEC.Data[7279] := 34.75;
   Prof_FEC.Data[7280] := 37.817;
   Prof_FEC.Data[7281] := 38.225;
   Prof_FEC.Data[7282] := 38.218;
   Prof_FEC.Data[7283] := 32.84;
   Prof_FEC.Data[7284] := 33.539;
   Prof_FEC.Data[7285] := 33.86;
   Prof_FEC.Data[7286] := 34.415;
   Prof_FEC.Data[7287] := 37.645;
   Prof_FEC.Data[7288] := 35.842;
   Prof_FEC.Data[7289] := 37.331;
   Prof_FEC.Data[7290] := 36.35;
   Prof_FEC.Data[7291] := 39.254;
   Prof_FEC.Data[7292] := 33.959;
   Prof_FEC.Data[7293] := 37.469;
   Prof_FEC.Data[7294] := 37.644;
   Prof_FEC.Data[7295] := 36.642;
   Prof_FEC.Data[7296] := 41.662;
   Prof_FEC.Data[7297] := 40.196;
   Prof_FEC.Data[7298] := 40.504;
   Prof_FEC.Data[7299] := 39.969;
   Prof_FEC.Data[7300] := 37.944;
   Prof_FEC.Data[7301] := 36.258;
   Prof_FEC.Data[7302] := 37.951;
   Prof_FEC.Data[7303] := 36.851;
   Prof_FEC.Data[7304] := 41.255;
   Prof_FEC.Data[7305] := 40.34;
   Prof_FEC.Data[7306] := 42.198;
   Prof_FEC.Data[7307] := 40.471;
   Prof_FEC.Data[7308] := 39.843;
   Prof_FEC.Data[7309] := 37.705;
   Prof_FEC.Data[7310] := 39.31;
   Prof_FEC.Data[7311] := 37.784;
   Prof_FEC.Data[7312] := 36.963;
   Prof_FEC.Data[7313] := 38.536;
   Prof_FEC.Data[7314] := 37.769;
   Prof_FEC.Data[7315] := 41.685;
   Prof_FEC.Data[7316] := 336.42;
   Prof_FEC.Data[7317] := 378.35;
   Prof_FEC.Data[7318] := 425.07;
   Prof_FEC.Data[7319] := 427.95;
   Prof_FEC.Data[7320] := 443.6;
   Prof_FEC.Data[7321] := 475.96;
   Prof_FEC.Data[7322] := 444.6;
   Prof_FEC.Data[7323] := 492.28;
   Prof_FEC.Data[7324] := 418.59;
   Prof_FEC.Data[7325] := 504.99;
   Prof_FEC.Data[7326] := 474.98;
   Prof_FEC.Data[7327] := 506.53;
   Prof_FEC.Data[7328] := 561.7;
   Prof_FEC.Data[7329] := 635.06;
   Prof_FEC.Data[7330] := 748.69;
   Prof_FEC.Data[7331] := 632.81;
   Prof_FEC.Data[7332] := 673.11;
   Prof_FEC.Data[7333] := 720.8;
   Prof_FEC.Data[7334] := 720.12;
   Prof_FEC.Data[7335] := 802.61;
   Prof_FEC.Data[7336] := 786.79;
   Prof_FEC.Data[7337] := 826.02;
   Prof_FEC.Data[7338] := 766.59;
   Prof_FEC.Data[7339] := 768.3;
   Prof_FEC.Data[7340] := 672.58;
   Prof_FEC.Data[7341] := 752.5;
   Prof_FEC.Data[7342] := 621.79;
   Prof_FEC.Data[7343] := 654.86;
   Prof_FEC.Data[7344] := 610.49;
   Prof_FEC.Data[7345] := 729.25;
   Prof_FEC.Data[7346] := 718.67;
   Prof_FEC.Data[7347] := 666.44;
   Prof_FEC.Data[7348] := 759.95;
   Prof_FEC.Data[7349] := 704.39;
   Prof_FEC.Data[7350] := 762.67;
   Prof_FEC.Data[7351] := 735.02;
   Prof_FEC.Data[7352] := 746.49;
   Prof_FEC.Data[7353] := 795.26;
   Prof_FEC.Data[7354] := 754.75;
   Prof_FEC.Data[7355] := 790.19;
   Prof_FEC.Data[7356] := 806.1;
   Prof_FEC.Data[7357] := 734.64;
   Prof_FEC.Data[7358] := 750.85;
   Prof_FEC.Data[7359] := 553.01;
   Prof_FEC.Data[7360] := 360.82;
   Prof_FEC.Data[7361] := 225.24;
   Prof_FEC.Data[7362] := 195.02;
   Prof_FEC.Data[7363] := 150.2;
   Prof_FEC.Data[7364] := 124.53;
   Prof_FEC.Data[7365] := 90.95;
   Prof_FEC.Data[7366] := 97.39;
   Prof_FEC.Data[7367] := 119.08;
   Prof_FEC.Data[7368] := 228.41;
   Prof_FEC.Data[7369] := 240.09;
   Prof_FEC.Data[7370] := 271.95;
   Prof_FEC.Data[7371] := 275.09;
   Prof_FEC.Data[7372] := 39.465;
   Prof_FEC.Data[7373] := 36.443;
   Prof_FEC.Data[7374] := 38.863;
   Prof_FEC.Data[7375] := 39.838;
   Prof_FEC.Data[7376] := 38.915;
   Prof_FEC.Data[7377] := 38.422;
   Prof_FEC.Data[7378] := 38.594;
   Prof_FEC.Data[7379] := 40.715;
   Prof_FEC.Data[7380] := 38.91;
   Prof_FEC.Data[7381] := 37.991;
   Prof_FEC.Data[7382] := 36.456;
   Prof_FEC.Data[7383] := 38.83;
   Prof_FEC.Data[7384] := 40.333;
   Prof_FEC.Data[7385] := 39.823;
   Prof_FEC.Data[7386] := 37.965;
   Prof_FEC.Data[7387] := 38.05;
   Prof_FEC.Data[7388] := 35.067;
   Prof_FEC.Data[7389] := 36.412;
   Prof_FEC.Data[7390] := 35.822;
   Prof_FEC.Data[7391] := 36.406;
   Prof_FEC.Data[7392] := 35.919;
   Prof_FEC.Data[7393] := 36.053;
   Prof_FEC.Data[7394] := 37.48;
   Prof_FEC.Data[7395] := 35.577;
   Prof_FEC.Data[7396] := 34.154;
   Prof_FEC.Data[7397] := 35.81;
   Prof_FEC.Data[7398] := 35.885;
   Prof_FEC.Data[7399] := 35.329;
   Prof_FEC.Data[7400] := 37.745;
   Prof_FEC.Data[7401] := 39.709;
   Prof_FEC.Data[7402] := 39.496;
   Prof_FEC.Data[7403] := 39.018;
   Prof_FEC.Data[7404] := 38.077;
   Prof_FEC.Data[7405] := 37.931;
   Prof_FEC.Data[7406] := 37.659;
   Prof_FEC.Data[7407] := 39.177;
   Prof_FEC.Data[7408] := 37.819;
   Prof_FEC.Data[7409] := 39.215;
   Prof_FEC.Data[7410] := 43.232;
   Prof_FEC.Data[7411] := 48.246;
   Prof_FEC.Data[7412] := 340.03;
   Prof_FEC.Data[7413] := 412.2;
   Prof_FEC.Data[7414] := 450.01;
   Prof_FEC.Data[7415] := 508.18;
   Prof_FEC.Data[7416] := 527.1;
   Prof_FEC.Data[7417] := 490.93;
   Prof_FEC.Data[7418] := 557.44;
   Prof_FEC.Data[7419] := 525.98;
   Prof_FEC.Data[7420] := 576.59;
   Prof_FEC.Data[7421] := 534.61;
   Prof_FEC.Data[7422] := 621.05;
   Prof_FEC.Data[7423] := 630.2;
   Prof_FEC.Data[7424] := 611.92;
   Prof_FEC.Data[7425] := 592.99;
   Prof_FEC.Data[7426] := 647.6;
   Prof_FEC.Data[7427] := 679.66;
   Prof_FEC.Data[7428] := 709.93;
   Prof_FEC.Data[7429] := 650.29;
   Prof_FEC.Data[7430] := 655.7;
   Prof_FEC.Data[7431] := 653.58;
   Prof_FEC.Data[7432] := 680.27;
   Prof_FEC.Data[7433] := 807.21;
   Prof_FEC.Data[7434] := 666.54;
   Prof_FEC.Data[7435] := 693.42;
   Prof_FEC.Data[7436] := 704.72;
   Prof_FEC.Data[7437] := 783.04;
   Prof_FEC.Data[7438] := 753.1;
   Prof_FEC.Data[7439] := 746.76;
   Prof_FEC.Data[7440] := 765.85;
   Prof_FEC.Data[7441] := 723.78;
   Prof_FEC.Data[7442] := 781.95;
   Prof_FEC.Data[7443] := 779.99;
   Prof_FEC.Data[7444] := 784.66;
   Prof_FEC.Data[7445] := 750.24;
   Prof_FEC.Data[7446] := 779.0;
   Prof_FEC.Data[7447] := 722.69;
   Prof_FEC.Data[7448] := 740.93;
   Prof_FEC.Data[7449] := 730.97;
   Prof_FEC.Data[7450] := 785.78;
   Prof_FEC.Data[7451] := 728.12;
   Prof_FEC.Data[7452] := 823.65;
   Prof_FEC.Data[7453] := 842.84;
   Prof_FEC.Data[7454] := 679.24;
   Prof_FEC.Data[7455] := 593.48;
   Prof_FEC.Data[7456] := 329.64;
   Prof_FEC.Data[7457] := 213.07;
   Prof_FEC.Data[7458] := 167.24;
   Prof_FEC.Data[7459] := 147.34;
   Prof_FEC.Data[7460] := 105.8;
   Prof_FEC.Data[7461] := 83.88;
   Prof_FEC.Data[7462] := 87.75;
   Prof_FEC.Data[7463] := 120.73;
   Prof_FEC.Data[7464] := 206.67;
   Prof_FEC.Data[7465] := 257.15;
   Prof_FEC.Data[7466] := 242.65;
   Prof_FEC.Data[7467] := 280.62;
   Prof_FEC.Data[7468] := 40.514;
   Prof_FEC.Data[7469] := 40.666;
   Prof_FEC.Data[7470] := 37.134;
   Prof_FEC.Data[7471] := 38.624;
   Prof_FEC.Data[7472] := 41.603;
   Prof_FEC.Data[7473] := 40.096;
   Prof_FEC.Data[7474] := 39.97;
   Prof_FEC.Data[7475] := 37.903;
   Prof_FEC.Data[7476] := 37.689;
   Prof_FEC.Data[7477] := 38.741;
   Prof_FEC.Data[7478] := 36.228;
   Prof_FEC.Data[7479] := 38.952;
   Prof_FEC.Data[7480] := 39.352;
   Prof_FEC.Data[7481] := 40.52;
   Prof_FEC.Data[7482] := 39.195;
   Prof_FEC.Data[7483] := 40.455;
   Prof_FEC.Data[7484] := 39.142;
   Prof_FEC.Data[7485] := 38.035;
   Prof_FEC.Data[7486] := 38.427;
   Prof_FEC.Data[7487] := 40.141;
   Prof_FEC.Data[7488] := 40.949;
   Prof_FEC.Data[7489] := 39.215;
   Prof_FEC.Data[7490] := 41.068;
   Prof_FEC.Data[7491] := 41.255;
   Prof_FEC.Data[7492] := 41.492;
   Prof_FEC.Data[7493] := 38.657;
   Prof_FEC.Data[7494] := 39.533;
   Prof_FEC.Data[7495] := 39.496;
   Prof_FEC.Data[7496] := 41.862;
   Prof_FEC.Data[7497] := 40.674;
   Prof_FEC.Data[7498] := 40.631;
   Prof_FEC.Data[7499] := 40.511;
   Prof_FEC.Data[7500] := 38.106;
   Prof_FEC.Data[7501] := 39.586;
   Prof_FEC.Data[7502] := 36.077;
   Prof_FEC.Data[7503] := 37.765;
   Prof_FEC.Data[7504] := 34.239;
   Prof_FEC.Data[7505] := 37.063;
   Prof_FEC.Data[7506] := 38.658;
   Prof_FEC.Data[7507] := 42.867;
   Prof_FEC.Data[7508] := 332.2;
   Prof_FEC.Data[7509] := 376.37;
   Prof_FEC.Data[7510] := 417.81;
   Prof_FEC.Data[7511] := 434.62;
   Prof_FEC.Data[7512] := 437.65;
   Prof_FEC.Data[7513] := 388.54;
   Prof_FEC.Data[7514] := 436.62;
   Prof_FEC.Data[7515] := 414.28;
   Prof_FEC.Data[7516] := 461.82;
   Prof_FEC.Data[7517] := 497.92;
   Prof_FEC.Data[7518] := 561.58;
   Prof_FEC.Data[7519] := 592.47;
   Prof_FEC.Data[7520] := 610.84;
   Prof_FEC.Data[7521] := 640.14;
   Prof_FEC.Data[7522] := 689.03;
   Prof_FEC.Data[7523] := 650.14;
   Prof_FEC.Data[7524] := 648.66;
   Prof_FEC.Data[7525] := 685.26;
   Prof_FEC.Data[7526] := 683.29;
   Prof_FEC.Data[7527] := 678.97;
   Prof_FEC.Data[7528] := 700.19;
   Prof_FEC.Data[7529] := 704.94;
   Prof_FEC.Data[7530] := 737.32;
   Prof_FEC.Data[7531] := 701.5;
   Prof_FEC.Data[7532] := 644.23;
   Prof_FEC.Data[7533] := 632.21;
   Prof_FEC.Data[7534] := 621.37;
   Prof_FEC.Data[7535] := 643.14;
   Prof_FEC.Data[7536] := 731.01;
   Prof_FEC.Data[7537] := 799.19;
   Prof_FEC.Data[7538] := 781.81;
   Prof_FEC.Data[7539] := 780.72;
   Prof_FEC.Data[7540] := 802.93;
   Prof_FEC.Data[7541] := 740.15;
   Prof_FEC.Data[7542] := 795.59;
   Prof_FEC.Data[7543] := 759.05;
   Prof_FEC.Data[7544] := 721.72;
   Prof_FEC.Data[7545] := 788.09;
   Prof_FEC.Data[7546] := 742.39;
   Prof_FEC.Data[7547] := 710.3;
   Prof_FEC.Data[7548] := 765.6;
   Prof_FEC.Data[7549] := 768.46;
   Prof_FEC.Data[7550] := 721.74;
   Prof_FEC.Data[7551] := 586.42;
   Prof_FEC.Data[7552] := 324.52;
   Prof_FEC.Data[7553] := 240.86;
   Prof_FEC.Data[7554] := 167.76;
   Prof_FEC.Data[7555] := 147.65;
   Prof_FEC.Data[7556] := 106.91;
   Prof_FEC.Data[7557] := 93.62;
   Prof_FEC.Data[7558] := 99.33;
   Prof_FEC.Data[7559] := 131.47;
   Prof_FEC.Data[7560] := 239.58;
   Prof_FEC.Data[7561] := 259.32;
   Prof_FEC.Data[7562] := 282.13;
   Prof_FEC.Data[7563] := 266.26;
   Prof_FEC.Data[7564] := 41.547;
   Prof_FEC.Data[7565] := 40.768;
   Prof_FEC.Data[7566] := 41.1;
   Prof_FEC.Data[7567] := 41.841;
   Prof_FEC.Data[7568] := 40.791;
   Prof_FEC.Data[7569] := 41.154;
   Prof_FEC.Data[7570] := 39.25;
   Prof_FEC.Data[7571] := 40.102;
   Prof_FEC.Data[7572] := 39.062;
   Prof_FEC.Data[7573] := 36.33;
   Prof_FEC.Data[7574] := 37.004;
   Prof_FEC.Data[7575] := 37.701;
   Prof_FEC.Data[7576] := 40.707;
   Prof_FEC.Data[7577] := 38.465;
   Prof_FEC.Data[7578] := 39.001;
   Prof_FEC.Data[7579] := 41.677;
   Prof_FEC.Data[7580] := 36.0;
   Prof_FEC.Data[7581] := 38.76;
   Prof_FEC.Data[7582] := 37.339;
   Prof_FEC.Data[7583] := 39.361;
   Prof_FEC.Data[7584] := 40.831;
   Prof_FEC.Data[7585] := 39.834;
   Prof_FEC.Data[7586] := 40.979;
   Prof_FEC.Data[7587] := 38.855;
   Prof_FEC.Data[7588] := 38.38;
   Prof_FEC.Data[7589] := 38.033;
   Prof_FEC.Data[7590] := 39.252;
   Prof_FEC.Data[7591] := 40.684;
   Prof_FEC.Data[7592] := 42.278;
   Prof_FEC.Data[7593] := 40.284;
   Prof_FEC.Data[7594] := 41.916;
   Prof_FEC.Data[7595] := 39.613;
   Prof_FEC.Data[7596] := 36.886;
   Prof_FEC.Data[7597] := 37.568;
   Prof_FEC.Data[7598] := 37.254;
   Prof_FEC.Data[7599] := 35.59;
   Prof_FEC.Data[7600] := 33.779;
   Prof_FEC.Data[7601] := 34.016;
   Prof_FEC.Data[7602] := 36.434;
   Prof_FEC.Data[7603] := 38.516;
   Prof_FEC.Data[7604] := 335.99;
   Prof_FEC.Data[7605] := 304.4;
   Prof_FEC.Data[7606] := 392.57;
   Prof_FEC.Data[7607] := 418.88;
   Prof_FEC.Data[7608] := 379.83;
   Prof_FEC.Data[7609] := 416.95;
   Prof_FEC.Data[7610] := 417.59;
   Prof_FEC.Data[7611] := 459.17;
   Prof_FEC.Data[7612] := 495.27;
   Prof_FEC.Data[7613] := 537.2;
   Prof_FEC.Data[7614] := 521.92;
   Prof_FEC.Data[7615] := 537.02;
   Prof_FEC.Data[7616] := 594.82;
   Prof_FEC.Data[7617] := 577.3;
   Prof_FEC.Data[7618] := 603.49;
   Prof_FEC.Data[7619] := 656.76;
   Prof_FEC.Data[7620] := 660.57;
   Prof_FEC.Data[7621] := 684.36;
   Prof_FEC.Data[7622] := 793.29;
   Prof_FEC.Data[7623] := 723.01;
   Prof_FEC.Data[7624] := 770.68;
   Prof_FEC.Data[7625] := 718.4;
   Prof_FEC.Data[7626] := 703.34;
   Prof_FEC.Data[7627] := 654.37;
   Prof_FEC.Data[7628] := 602.49;
   Prof_FEC.Data[7629] := 613.98;
   Prof_FEC.Data[7630] := 565.79;
   Prof_FEC.Data[7631] := 545.27;
   Prof_FEC.Data[7632] := 586.14;
   Prof_FEC.Data[7633] := 649.87;
   Prof_FEC.Data[7634] := 583.78;
   Prof_FEC.Data[7635] := 635.24;
   Prof_FEC.Data[7636] := 631.88;
   Prof_FEC.Data[7637] := 582.62;
   Prof_FEC.Data[7638] := 634.88;
   Prof_FEC.Data[7639] := 601.99;
   Prof_FEC.Data[7640] := 633.44;
   Prof_FEC.Data[7641] := 621.58;
   Prof_FEC.Data[7642] := 622.87;
   Prof_FEC.Data[7643] := 597.48;
   Prof_FEC.Data[7644] := 634.07;
   Prof_FEC.Data[7645] := 694.23;
   Prof_FEC.Data[7646] := 748.59;
   Prof_FEC.Data[7647] := 500.55;
   Prof_FEC.Data[7648] := 291.24;
   Prof_FEC.Data[7649] := 205.77;
   Prof_FEC.Data[7650] := 146.14;
   Prof_FEC.Data[7651] := 135.23;
   Prof_FEC.Data[7652] := 111.13;
   Prof_FEC.Data[7653] := 93.13;
   Prof_FEC.Data[7654] := 93.47;
   Prof_FEC.Data[7655] := 121.82;
   Prof_FEC.Data[7656] := 195.44;
   Prof_FEC.Data[7657] := 230.53;
   Prof_FEC.Data[7658] := 264.34;
   Prof_FEC.Data[7659] := 238.27;
   Prof_FEC.Data[7660] := 39.043;
   Prof_FEC.Data[7661] := 36.481;
   Prof_FEC.Data[7662] := 39.071;
   Prof_FEC.Data[7663] := 37.702;
   Prof_FEC.Data[7664] := 40.46;
   Prof_FEC.Data[7665] := 39.95;
   Prof_FEC.Data[7666] := 41.594;
   Prof_FEC.Data[7667] := 39.557;
   Prof_FEC.Data[7668] := 38.159;
   Prof_FEC.Data[7669] := 38.937;
   Prof_FEC.Data[7670] := 36.935;
   Prof_FEC.Data[7671] := 40.03;
   Prof_FEC.Data[7672] := 40.568;
   Prof_FEC.Data[7673] := 40.859;
   Prof_FEC.Data[7674] := 44.084;
   Prof_FEC.Data[7675] := 41.64;
   Prof_FEC.Data[7676] := 37.833;
   Prof_FEC.Data[7677] := 40.578;
   Prof_FEC.Data[7678] := 38.093;
   Prof_FEC.Data[7679] := 40.191;
   Prof_FEC.Data[7680] := 40.509;
   Prof_FEC.Data[7681] := 37.185;
   Prof_FEC.Data[7682] := 41.031;
   Prof_FEC.Data[7683] := 39.722;
   Prof_FEC.Data[7684] := 38.497;
   Prof_FEC.Data[7685] := 37.751;
   Prof_FEC.Data[7686] := 38.696;
   Prof_FEC.Data[7687] := 37.076;
   Prof_FEC.Data[7688] := 40.397;
   Prof_FEC.Data[7689] := 37.349;
   Prof_FEC.Data[7690] := 39.803;
   Prof_FEC.Data[7691] := 38.737;
   Prof_FEC.Data[7692] := 37.377;
   Prof_FEC.Data[7693] := 36.419;
   Prof_FEC.Data[7694] := 35.564;
   Prof_FEC.Data[7695] := 36.816;
   Prof_FEC.Data[7696] := 37.074;
   Prof_FEC.Data[7697] := 38.239;
   Prof_FEC.Data[7698] := 37.615;
   Prof_FEC.Data[7699] := 37.18;
   Prof_FEC.Data[7700] := 224.23;
   Prof_FEC.Data[7701] := 182.52;
   Prof_FEC.Data[7702] := 217.42;
   Prof_FEC.Data[7703] := 208.8;
   Prof_FEC.Data[7704] := 234.0;
   Prof_FEC.Data[7705] := 245.69;
   Prof_FEC.Data[7706] := 271.4;
   Prof_FEC.Data[7707] := 310.44;
   Prof_FEC.Data[7708] := 286.19;
   Prof_FEC.Data[7709] := 281.09;
   Prof_FEC.Data[7710] := 334.91;
   Prof_FEC.Data[7711] := 308.25;
   Prof_FEC.Data[7712] := 338.3;
   Prof_FEC.Data[7713] := 356.72;
   Prof_FEC.Data[7714] := 364.0;
   Prof_FEC.Data[7715] := 398.07;
   Prof_FEC.Data[7716] := 406.77;
   Prof_FEC.Data[7717] := 422.21;
   Prof_FEC.Data[7718] := 429.88;
   Prof_FEC.Data[7719] := 405.24;
   Prof_FEC.Data[7720] := 457.44;
   Prof_FEC.Data[7721] := 434.43;
   Prof_FEC.Data[7722] := 414.75;
   Prof_FEC.Data[7723] := 353.77;
   Prof_FEC.Data[7724] := 294.66;
   Prof_FEC.Data[7725] := 302.55;
   Prof_FEC.Data[7726] := 293.61;
   Prof_FEC.Data[7727] := 273.0;
   Prof_FEC.Data[7728] := 304.56;
   Prof_FEC.Data[7729] := 295.35;
   Prof_FEC.Data[7730] := 285.0;
   Prof_FEC.Data[7731] := 266.08;
   Prof_FEC.Data[7732] := 272.21;
   Prof_FEC.Data[7733] := 285.99;
   Prof_FEC.Data[7734] := 300.28;
   Prof_FEC.Data[7735] := 303.17;
   Prof_FEC.Data[7736] := 307.71;
   Prof_FEC.Data[7737] := 304.22;
   Prof_FEC.Data[7738] := 294.83;
   Prof_FEC.Data[7739] := 218.74;
   Prof_FEC.Data[7740] := 144.72;
   Prof_FEC.Data[7741] := 103.12;
   Prof_FEC.Data[7742] := 80.14;
   Prof_FEC.Data[7743] := 75.28;
   Prof_FEC.Data[7744] := 89.68;
   Prof_FEC.Data[7745] := 91.93;
   Prof_FEC.Data[7746] := 88.21;
   Prof_FEC.Data[7747] := 94.12;
   Prof_FEC.Data[7748] := 93.29;
   Prof_FEC.Data[7749] := 97.86;
   Prof_FEC.Data[7750] := 105.64;
   Prof_FEC.Data[7751] := 154.93;
   Prof_FEC.Data[7752] := 164.74;
   Prof_FEC.Data[7753] := 200.11;
   Prof_FEC.Data[7754] := 237.73;
   Prof_FEC.Data[7755] := 236.91;
   Prof_FEC.Data[7756] := 39.125;
   Prof_FEC.Data[7757] := 40.242;
   Prof_FEC.Data[7758] := 41.14;
   Prof_FEC.Data[7759] := 38.696;
   Prof_FEC.Data[7760] := 38.027;
   Prof_FEC.Data[7761] := 33.638;
   Prof_FEC.Data[7762] := 34.131;
   Prof_FEC.Data[7763] := 35.772;
   Prof_FEC.Data[7764] := 38.755;
   Prof_FEC.Data[7765] := 35.307;
   Prof_FEC.Data[7766] := 35.464;
   Prof_FEC.Data[7767] := 36.856;
   Prof_FEC.Data[7768] := 36.57;
   Prof_FEC.Data[7769] := 35.455;
   Prof_FEC.Data[7770] := 35.575;
   Prof_FEC.Data[7771] := 36.98;
   Prof_FEC.Data[7772] := 38.359;
   Prof_FEC.Data[7773] := 37.828;
   Prof_FEC.Data[7774] := 38.9;
   Prof_FEC.Data[7775] := 37.14;
   Prof_FEC.Data[7776] := 36.647;
   Prof_FEC.Data[7777] := 36.455;
   Prof_FEC.Data[7778] := 34.957;
   Prof_FEC.Data[7779] := 36.962;
   Prof_FEC.Data[7780] := 36.264;
   Prof_FEC.Data[7781] := 38.303;
   Prof_FEC.Data[7782] := 38.018;
   Prof_FEC.Data[7783] := 38.787;
   Prof_FEC.Data[7784] := 38.188;
   Prof_FEC.Data[7785] := 37.398;
   Prof_FEC.Data[7786] := 36.257;
   Prof_FEC.Data[7787] := 37.307;
   Prof_FEC.Data[7788] := 38.834;
   Prof_FEC.Data[7789] := 42.187;
   Prof_FEC.Data[7790] := 39.275;
   Prof_FEC.Data[7791] := 37.488;
   Prof_FEC.Data[7792] := 34.589;
   Prof_FEC.Data[7793] := 36.53;
   Prof_FEC.Data[7794] := 37.429;
   Prof_FEC.Data[7795] := 36.17;
   Prof_FEC.Data[7796] := 236.05;
   Prof_FEC.Data[7797] := 237.86;
   Prof_FEC.Data[7798] := 227.9;
   Prof_FEC.Data[7799] := 218.89;
   Prof_FEC.Data[7800] := 180.6;
   Prof_FEC.Data[7801] := 137.16;
   Prof_FEC.Data[7802] := 131.42;
   Prof_FEC.Data[7803] := 123.52;
   Prof_FEC.Data[7804] := 114.59;
   Prof_FEC.Data[7805] := 116.78;
   Prof_FEC.Data[7806] := 109.02;
   Prof_FEC.Data[7807] := 126.96;
   Prof_FEC.Data[7808] := 129.85;
   Prof_FEC.Data[7809] := 114.98;
   Prof_FEC.Data[7810] := 111.69;
   Prof_FEC.Data[7811] := 114.36;
   Prof_FEC.Data[7812] := 125.31;
   Prof_FEC.Data[7813] := 145.83;
   Prof_FEC.Data[7814] := 136.67;
   Prof_FEC.Data[7815] := 137.52;
   Prof_FEC.Data[7816] := 121.57;
   Prof_FEC.Data[7817] := 129.88;
   Prof_FEC.Data[7818] := 121.1;
   Prof_FEC.Data[7819] := 120.62;
   Prof_FEC.Data[7820] := 144.79;
   Prof_FEC.Data[7821] := 131.58;
   Prof_FEC.Data[7822] := 138.17;
   Prof_FEC.Data[7823] := 137.86;
   Prof_FEC.Data[7824] := 119.15;
   Prof_FEC.Data[7825] := 109.65;
   Prof_FEC.Data[7826] := 114.37;
   Prof_FEC.Data[7827] := 112.38;
   Prof_FEC.Data[7828] := 139.48;
   Prof_FEC.Data[7829] := 146.95;
   Prof_FEC.Data[7830] := 147.62;
   Prof_FEC.Data[7831] := 132.26;
   Prof_FEC.Data[7832] := 146.92;
   Prof_FEC.Data[7833] := 126.45;
   Prof_FEC.Data[7834] := 130.09;
   Prof_FEC.Data[7835] := 124.75;
   Prof_FEC.Data[7836] := 136.72;
   Prof_FEC.Data[7837] := 151.58;
   Prof_FEC.Data[7838] := 139.95;
   Prof_FEC.Data[7839] := 131.48;
   Prof_FEC.Data[7840] := 122.36;
   Prof_FEC.Data[7841] := 123.93;
   Prof_FEC.Data[7842] := 112.2;
   Prof_FEC.Data[7843] := 117.94;
   Prof_FEC.Data[7844] := 121.51;
   Prof_FEC.Data[7845] := 124.63;
   Prof_FEC.Data[7846] := 141.59;
   Prof_FEC.Data[7847] := 176.8;
   Prof_FEC.Data[7848] := 206.93;
   Prof_FEC.Data[7849] := 223.66;
   Prof_FEC.Data[7850] := 227.34;
   Prof_FEC.Data[7851] := 243.91;
   Prof_FEC.Data[7852] := 41.164;
   Prof_FEC.Data[7853] := 45.574;
   Prof_FEC.Data[7854] := 43.955;
   Prof_FEC.Data[7855] := 44.214;
   Prof_FEC.Data[7856] := 41.107;
   Prof_FEC.Data[7857] := 38.803;
   Prof_FEC.Data[7858] := 40.838;
   Prof_FEC.Data[7859] := 40.29;
   Prof_FEC.Data[7860] := 43.656;
   Prof_FEC.Data[7861] := 41.745;
   Prof_FEC.Data[7862] := 39.977;
   Prof_FEC.Data[7863] := 40.914;
   Prof_FEC.Data[7864] := 38.535;
   Prof_FEC.Data[7865] := 38.606;
   Prof_FEC.Data[7866] := 35.907;
   Prof_FEC.Data[7867] := 36.845;
   Prof_FEC.Data[7868] := 39.165;
   Prof_FEC.Data[7869] := 38.546;
   Prof_FEC.Data[7870] := 40.647;
   Prof_FEC.Data[7871] := 40.367;
   Prof_FEC.Data[7872] := 40.244;
   Prof_FEC.Data[7873] := 37.594;
   Prof_FEC.Data[7874] := 37.255;
   Prof_FEC.Data[7875] := 36.185;
   Prof_FEC.Data[7876] := 38.218;
   Prof_FEC.Data[7877] := 36.94;
   Prof_FEC.Data[7878] := 38.157;
   Prof_FEC.Data[7879] := 37.315;
   Prof_FEC.Data[7880] := 36.431;
   Prof_FEC.Data[7881] := 36.131;
   Prof_FEC.Data[7882] := 36.748;
   Prof_FEC.Data[7883] := 38.317;
   Prof_FEC.Data[7884] := 33.749;
   Prof_FEC.Data[7885] := 36.936;
   Prof_FEC.Data[7886] := 38.394;
   Prof_FEC.Data[7887] := 36.215;
   Prof_FEC.Data[7888] := 35.455;
   Prof_FEC.Data[7889] := 35.564;
   Prof_FEC.Data[7890] := 34.277;
   Prof_FEC.Data[7891] := 36.35;
   Prof_FEC.Data[7892] := 294.36;
   Prof_FEC.Data[7893] := 317.77;
   Prof_FEC.Data[7894] := 348.52;
   Prof_FEC.Data[7895] := 363.49;
   Prof_FEC.Data[7896] := 372.84;
   Prof_FEC.Data[7897] := 369.69;
   Prof_FEC.Data[7898] := 415.16;
   Prof_FEC.Data[7899] := 449.48;
   Prof_FEC.Data[7900] := 481.36;
   Prof_FEC.Data[7901] := 555.58;
   Prof_FEC.Data[7902] := 526.88;
   Prof_FEC.Data[7903] := 546.84;
   Prof_FEC.Data[7904] := 550.7;
   Prof_FEC.Data[7905] := 525.77;
   Prof_FEC.Data[7906] := 615.35;
   Prof_FEC.Data[7907] := 609.06;
   Prof_FEC.Data[7908] := 631.06;
   Prof_FEC.Data[7909] := 643.89;
   Prof_FEC.Data[7910] := 611.6;
   Prof_FEC.Data[7911] := 636.42;
   Prof_FEC.Data[7912] := 657.97;
   Prof_FEC.Data[7913] := 752.98;
   Prof_FEC.Data[7914] := 674.23;
   Prof_FEC.Data[7915] := 640.57;
   Prof_FEC.Data[7916] := 580.8;
   Prof_FEC.Data[7917] := 613.26;
   Prof_FEC.Data[7918] := 581.0;
   Prof_FEC.Data[7919] := 623.05;
   Prof_FEC.Data[7920] := 693.83;
   Prof_FEC.Data[7921] := 710.9;
   Prof_FEC.Data[7922] := 739.42;
   Prof_FEC.Data[7923] := 705.58;
   Prof_FEC.Data[7924] := 650.67;
   Prof_FEC.Data[7925] := 660.51;
   Prof_FEC.Data[7926] := 648.39;
   Prof_FEC.Data[7927] := 646.16;
   Prof_FEC.Data[7928] := 567.23;
   Prof_FEC.Data[7929] := 616.9;
   Prof_FEC.Data[7930] := 611.89;
   Prof_FEC.Data[7931] := 624.87;
   Prof_FEC.Data[7932] := 705.38;
   Prof_FEC.Data[7933] := 703.64;
   Prof_FEC.Data[7934] := 707.9;
   Prof_FEC.Data[7935] := 617.65;
   Prof_FEC.Data[7936] := 353.74;
   Prof_FEC.Data[7937] := 240.12;
   Prof_FEC.Data[7938] := 189.46;
   Prof_FEC.Data[7939] := 161.54;
   Prof_FEC.Data[7940] := 123.08;
   Prof_FEC.Data[7941] := 113.68;
   Prof_FEC.Data[7942] := 115.78;
   Prof_FEC.Data[7943] := 123.65;
   Prof_FEC.Data[7944] := 229.55;
   Prof_FEC.Data[7945] := 237.9;
   Prof_FEC.Data[7946] := 251.59;
   Prof_FEC.Data[7947] := 255.8;
   Prof_FEC.Data[7948] := 40.26;
   Prof_FEC.Data[7949] := 37.918;
   Prof_FEC.Data[7950] := 37.914;
   Prof_FEC.Data[7951] := 39.097;
   Prof_FEC.Data[7952] := 41.255;
   Prof_FEC.Data[7953] := 41.5;
   Prof_FEC.Data[7954] := 40.119;
   Prof_FEC.Data[7955] := 38.425;
   Prof_FEC.Data[7956] := 35.738;
   Prof_FEC.Data[7957] := 39.833;
   Prof_FEC.Data[7958] := 36.7;
   Prof_FEC.Data[7959] := 37.574;
   Prof_FEC.Data[7960] := 38.951;
   Prof_FEC.Data[7961] := 39.196;
   Prof_FEC.Data[7962] := 40.034;
   Prof_FEC.Data[7963] := 41.039;
   Prof_FEC.Data[7964] := 40.562;
   Prof_FEC.Data[7965] := 40.896;
   Prof_FEC.Data[7966] := 41.183;
   Prof_FEC.Data[7967] := 39.083;
   Prof_FEC.Data[7968] := 41.112;
   Prof_FEC.Data[7969] := 42.98;
   Prof_FEC.Data[7970] := 41.46;
   Prof_FEC.Data[7971] := 40.185;
   Prof_FEC.Data[7972] := 39.799;
   Prof_FEC.Data[7973] := 39.77;
   Prof_FEC.Data[7974] := 38.476;
   Prof_FEC.Data[7975] := 39.703;
   Prof_FEC.Data[7976] := 42.937;
   Prof_FEC.Data[7977] := 42.328;
   Prof_FEC.Data[7978] := 41.814;
   Prof_FEC.Data[7979] := 38.641;
   Prof_FEC.Data[7980] := 39.146;
   Prof_FEC.Data[7981] := 37.497;
   Prof_FEC.Data[7982] := 36.529;
   Prof_FEC.Data[7983] := 38.061;
   Prof_FEC.Data[7984] := 39.216;
   Prof_FEC.Data[7985] := 39.229;
   Prof_FEC.Data[7986] := 39.049;
   Prof_FEC.Data[7987] := 42.388;
   Prof_FEC.Data[7988] := 356.95;
   Prof_FEC.Data[7989] := 383.66;
   Prof_FEC.Data[7990] := 427.0;
   Prof_FEC.Data[7991] := 403.55;
   Prof_FEC.Data[7992] := 443.25;
   Prof_FEC.Data[7993] := 412.66;
   Prof_FEC.Data[7994] := 475.12;
   Prof_FEC.Data[7995] := 434.3;
   Prof_FEC.Data[7996] := 574.04;
   Prof_FEC.Data[7997] := 568.99;
   Prof_FEC.Data[7998] := 579.74;
   Prof_FEC.Data[7999] := 582.87;
   Prof_FEC.Data[8000] := 574.86;
   Prof_FEC.Data[8001] := 712.43;
   Prof_FEC.Data[8002] := 683.15;
   Prof_FEC.Data[8003] := 725.59;
   Prof_FEC.Data[8004] := 675.92;
   Prof_FEC.Data[8005] := 700.98;
   Prof_FEC.Data[8006] := 643.74;
   Prof_FEC.Data[8007] := 696.07;
   Prof_FEC.Data[8008] := 646.2;
   Prof_FEC.Data[8009] := 842.24;
   Prof_FEC.Data[8010] := 695.42;
   Prof_FEC.Data[8011] := 670.74;
   Prof_FEC.Data[8012] := 590.43;
   Prof_FEC.Data[8013] := 594.78;
   Prof_FEC.Data[8014] := 630.22;
   Prof_FEC.Data[8015] := 543.74;
   Prof_FEC.Data[8016] := 573.58;
   Prof_FEC.Data[8017] := 628.97;
   Prof_FEC.Data[8018] := 618.39;
   Prof_FEC.Data[8019] := 602.45;
   Prof_FEC.Data[8020] := 640.51;
   Prof_FEC.Data[8021] := 633.84;
   Prof_FEC.Data[8022] := 599.69;
   Prof_FEC.Data[8023] := 611.95;
   Prof_FEC.Data[8024] := 659.83;
   Prof_FEC.Data[8025] := 696.86;
   Prof_FEC.Data[8026] := 727.57;
   Prof_FEC.Data[8027] := 628.04;
   Prof_FEC.Data[8028] := 657.14;
   Prof_FEC.Data[8029] := 729.72;
   Prof_FEC.Data[8030] := 642.29;
   Prof_FEC.Data[8031] := 549.53;
   Prof_FEC.Data[8032] := 303.19;
   Prof_FEC.Data[8033] := 190.66;
   Prof_FEC.Data[8034] := 119.37;
   Prof_FEC.Data[8035] := 100.56;
   Prof_FEC.Data[8036] := 68.24;
   Prof_FEC.Data[8037] := 51.05;
   Prof_FEC.Data[8038] := 68.44;
   Prof_FEC.Data[8039] := 79.19;
   Prof_FEC.Data[8040] := 142.55;
   Prof_FEC.Data[8041] := 137.14;
   Prof_FEC.Data[8042] := 198.39;
   Prof_FEC.Data[8043] := 201.05;
   Prof_FEC.Data[8044] := 31.465;
   Prof_FEC.Data[8045] := 33.704;
   Prof_FEC.Data[8046] := 34.405;
   Prof_FEC.Data[8047] := 32.884;
   Prof_FEC.Data[8048] := 35.406;
   Prof_FEC.Data[8049] := 37.471;
   Prof_FEC.Data[8050] := 36.902;
   Prof_FEC.Data[8051] := 34.323;
   Prof_FEC.Data[8052] := 35.049;
   Prof_FEC.Data[8053] := 37.428;
   Prof_FEC.Data[8054] := 37.559;
   Prof_FEC.Data[8055] := 38.833;
   Prof_FEC.Data[8056] := 40.594;
   Prof_FEC.Data[8057] := 38.67;
   Prof_FEC.Data[8058] := 41.709;
   Prof_FEC.Data[8059] := 40.129;
   Prof_FEC.Data[8060] := 38.75;
   Prof_FEC.Data[8061] := 37.905;
   Prof_FEC.Data[8062] := 36.95;
   Prof_FEC.Data[8063] := 36.541;
   Prof_FEC.Data[8064] := 37.066;
   Prof_FEC.Data[8065] := 41.044;
   Prof_FEC.Data[8066] := 39.2;
   Prof_FEC.Data[8067] := 35.61;
   Prof_FEC.Data[8068] := 36.134;
   Prof_FEC.Data[8069] := 32.693;
   Prof_FEC.Data[8070] := 35.759;
   Prof_FEC.Data[8071] := 36.637;
   Prof_FEC.Data[8072] := 37.385;
   Prof_FEC.Data[8073] := 36.888;
   Prof_FEC.Data[8074] := 39.161;
   Prof_FEC.Data[8075] := 37.836;
   Prof_FEC.Data[8076] := 33.957;
   Prof_FEC.Data[8077] := 37.954;
   Prof_FEC.Data[8078] := 36.334;
   Prof_FEC.Data[8079] := 37.126;
   Prof_FEC.Data[8080] := 39.331;
   Prof_FEC.Data[8081] := 40.392;
   Prof_FEC.Data[8082] := 40.182;
   Prof_FEC.Data[8083] := 42.871;
   Prof_FEC.Data[8084] := 339.04;
   Prof_FEC.Data[8085] := 382.04;
   Prof_FEC.Data[8086] := 410.09;
   Prof_FEC.Data[8087] := 423.45;
   Prof_FEC.Data[8088] := 395.17;
   Prof_FEC.Data[8089] := 414.51;
   Prof_FEC.Data[8090] := 443.09;
   Prof_FEC.Data[8091] := 438.45;
   Prof_FEC.Data[8092] := 454.17;
   Prof_FEC.Data[8093] := 518.75;
   Prof_FEC.Data[8094] := 553.41;
   Prof_FEC.Data[8095] := 554.79;
   Prof_FEC.Data[8096] := 664.85;
   Prof_FEC.Data[8097] := 621.4;
   Prof_FEC.Data[8098] := 633.69;
   Prof_FEC.Data[8099] := 602.23;
   Prof_FEC.Data[8100] := 672.11;
   Prof_FEC.Data[8101] := 672.8;
   Prof_FEC.Data[8102] := 652.54;
   Prof_FEC.Data[8103] := 628.43;
   Prof_FEC.Data[8104] := 567.49;
   Prof_FEC.Data[8105] := 540.9;
   Prof_FEC.Data[8106] := 607.09;
   Prof_FEC.Data[8107] := 567.82;
   Prof_FEC.Data[8108] := 564.5;
   Prof_FEC.Data[8109] := 569.05;
   Prof_FEC.Data[8110] := 557.25;
   Prof_FEC.Data[8111] := 521.32;
   Prof_FEC.Data[8112] := 667.19;
   Prof_FEC.Data[8113] := 644.19;
   Prof_FEC.Data[8114] := 663.54;
   Prof_FEC.Data[8115] := 636.21;
   Prof_FEC.Data[8116] := 649.11;
   Prof_FEC.Data[8117] := 577.0;
   Prof_FEC.Data[8118] := 628.22;
   Prof_FEC.Data[8119] := 619.05;
   Prof_FEC.Data[8120] := 657.88;
   Prof_FEC.Data[8121] := 642.18;
   Prof_FEC.Data[8122] := 645.27;
   Prof_FEC.Data[8123] := 651.4;
   Prof_FEC.Data[8124] := 685.61;
   Prof_FEC.Data[8125] := 738.71;
   Prof_FEC.Data[8126] := 548.33;
   Prof_FEC.Data[8127] := 478.7;
   Prof_FEC.Data[8128] := 278.12;
   Prof_FEC.Data[8129] := 167.23;
   Prof_FEC.Data[8130] := 128.06;
   Prof_FEC.Data[8131] := 120.28;
   Prof_FEC.Data[8132] := 80.33;
   Prof_FEC.Data[8133] := 58.08;
   Prof_FEC.Data[8134] := 65.33;
   Prof_FEC.Data[8135] := 80.24;
   Prof_FEC.Data[8136] := 134.84;
   Prof_FEC.Data[8137] := 145.97;
   Prof_FEC.Data[8138] := 183.78;
   Prof_FEC.Data[8139] := 196.29;
   Prof_FEC.Data[8140] := 33.488;
   Prof_FEC.Data[8141] := 33.235;
   Prof_FEC.Data[8142] := 34.273;
   Prof_FEC.Data[8143] := 33.556;
   Prof_FEC.Data[8144] := 35.353;
   Prof_FEC.Data[8145] := 35.156;
   Prof_FEC.Data[8146] := 37.721;
   Prof_FEC.Data[8147] := 36.51;
   Prof_FEC.Data[8148] := 34.46;
   Prof_FEC.Data[8149] := 36.289;
   Prof_FEC.Data[8150] := 36.751;
   Prof_FEC.Data[8151] := 37.643;
   Prof_FEC.Data[8152] := 37.642;
   Prof_FEC.Data[8153] := 38.147;
   Prof_FEC.Data[8154] := 41.717;
   Prof_FEC.Data[8155] := 37.499;
   Prof_FEC.Data[8156] := 38.388;
   Prof_FEC.Data[8157] := 38.031;
   Prof_FEC.Data[8158] := 37.422;
   Prof_FEC.Data[8159] := 36.964;
   Prof_FEC.Data[8160] := 42.666;
   Prof_FEC.Data[8161] := 41.232;
   Prof_FEC.Data[8162] := 41.387;
   Prof_FEC.Data[8163] := 41.556;
   Prof_FEC.Data[8164] := 39.69;
   Prof_FEC.Data[8165] := 37.528;
   Prof_FEC.Data[8166] := 36.845;
   Prof_FEC.Data[8167] := 40.682;
   Prof_FEC.Data[8168] := 39.759;
   Prof_FEC.Data[8169] := 41.845;
   Prof_FEC.Data[8170] := 43.777;
   Prof_FEC.Data[8171] := 40.177;
   Prof_FEC.Data[8172] := 36.81;
   Prof_FEC.Data[8173] := 36.916;
   Prof_FEC.Data[8174] := 38.027;
   Prof_FEC.Data[8175] := 38.115;
   Prof_FEC.Data[8176] := 39.079;
   Prof_FEC.Data[8177] := 38.708;
   Prof_FEC.Data[8178] := 37.383;
   Prof_FEC.Data[8179] := 46.836;
   Prof_FEC.Data[8180] := 326.93;
   Prof_FEC.Data[8181] := 385.36;
   Prof_FEC.Data[8182] := 418.04;
   Prof_FEC.Data[8183] := 408.57;
   Prof_FEC.Data[8184] := 404.75;
   Prof_FEC.Data[8185] := 412.01;
   Prof_FEC.Data[8186] := 425.73;
   Prof_FEC.Data[8187] := 459.78;
   Prof_FEC.Data[8188] := 447.81;
   Prof_FEC.Data[8189] := 578.22;
   Prof_FEC.Data[8190] := 538.09;
   Prof_FEC.Data[8191] := 629.99;
   Prof_FEC.Data[8192] := 581.96;
   Prof_FEC.Data[8193] := 607.13;
   Prof_FEC.Data[8194] := 668.57;
   Prof_FEC.Data[8195] := 622.16;
   Prof_FEC.Data[8196] := 636.06;
   Prof_FEC.Data[8197] := 670.34;
   Prof_FEC.Data[8198] := 648.57;
   Prof_FEC.Data[8199] := 603.47;
   Prof_FEC.Data[8200] := 611.41;
   Prof_FEC.Data[8201] := 550.22;
   Prof_FEC.Data[8202] := 616.31;
   Prof_FEC.Data[8203] := 623.23;
   Prof_FEC.Data[8204] := 555.19;
   Prof_FEC.Data[8205] := 568.24;
   Prof_FEC.Data[8206] := 583.24;
   Prof_FEC.Data[8207] := 661.89;
   Prof_FEC.Data[8208] := 640.43;
   Prof_FEC.Data[8209] := 648.32;
   Prof_FEC.Data[8210] := 663.08;
   Prof_FEC.Data[8211] := 651.73;
   Prof_FEC.Data[8212] := 642.23;
   Prof_FEC.Data[8213] := 694.44;
   Prof_FEC.Data[8214] := 676.12;
   Prof_FEC.Data[8215] := 749.53;
   Prof_FEC.Data[8216] := 731.88;
   Prof_FEC.Data[8217] := 773.44;
   Prof_FEC.Data[8218] := 753.7;
   Prof_FEC.Data[8219] := 698.73;
   Prof_FEC.Data[8220] := 801.99;
   Prof_FEC.Data[8221] := 761.02;
   Prof_FEC.Data[8222] := 724.45;
   Prof_FEC.Data[8223] := 602.65;
   Prof_FEC.Data[8224] := 301.99;
   Prof_FEC.Data[8225] := 194.1;
   Prof_FEC.Data[8226] := 133.57;
   Prof_FEC.Data[8227] := 113.14;
   Prof_FEC.Data[8228] := 85.79;
   Prof_FEC.Data[8229] := 71.46;
   Prof_FEC.Data[8230] := 68.26;
   Prof_FEC.Data[8231] := 99.1;
   Prof_FEC.Data[8232] := 174.15;
   Prof_FEC.Data[8233] := 198.57;
   Prof_FEC.Data[8234] := 209.34;
   Prof_FEC.Data[8235] := 228.34;
   Prof_FEC.Data[8236] := 38.17;
   Prof_FEC.Data[8237] := 39.136;
   Prof_FEC.Data[8238] := 37.265;
   Prof_FEC.Data[8239] := 38.564;
   Prof_FEC.Data[8240] := 37.998;
   Prof_FEC.Data[8241] := 38.232;
   Prof_FEC.Data[8242] := 37.622;
   Prof_FEC.Data[8243] := 38.082;
   Prof_FEC.Data[8244] := 37.489;
   Prof_FEC.Data[8245] := 34.913;
   Prof_FEC.Data[8246] := 36.065;
   Prof_FEC.Data[8247] := 36.828;
   Prof_FEC.Data[8248] := 34.984;
   Prof_FEC.Data[8249] := 37.465;
   Prof_FEC.Data[8250] := 37.485;
   Prof_FEC.Data[8251] := 36.792;
   Prof_FEC.Data[8252] := 35.377;
   Prof_FEC.Data[8253] := 35.906;
   Prof_FEC.Data[8254] := 36.837;
   Prof_FEC.Data[8255] := 39.485;
   Prof_FEC.Data[8256] := 38.128;
   Prof_FEC.Data[8257] := 37.919;
   Prof_FEC.Data[8258] := 36.893;
   Prof_FEC.Data[8259] := 37.368;
   Prof_FEC.Data[8260] := 36.47;
   Prof_FEC.Data[8261] := 37.671;
   Prof_FEC.Data[8262] := 35.255;
   Prof_FEC.Data[8263] := 36.979;
   Prof_FEC.Data[8264] := 36.243;
   Prof_FEC.Data[8265] := 41.015;
   Prof_FEC.Data[8266] := 39.576;
   Prof_FEC.Data[8267] := 40.556;
   Prof_FEC.Data[8268] := 37.06;
   Prof_FEC.Data[8269] := 38.161;
   Prof_FEC.Data[8270] := 38.193;
   Prof_FEC.Data[8271] := 36.126;
   Prof_FEC.Data[8272] := 33.95;
   Prof_FEC.Data[8273] := 35.968;
   Prof_FEC.Data[8274] := 38.233;
   Prof_FEC.Data[8275] := 41.701;
   Prof_FEC.Data[8276] := 330.44;
   Prof_FEC.Data[8277] := 371.91;
   Prof_FEC.Data[8278] := 388.56;
   Prof_FEC.Data[8279] := 427.35;
   Prof_FEC.Data[8280] := 372.05;
   Prof_FEC.Data[8281] := 352.33;
   Prof_FEC.Data[8282] := 415.79;
   Prof_FEC.Data[8283] := 474.41;
   Prof_FEC.Data[8284] := 529.5;
   Prof_FEC.Data[8285] := 592.28;
   Prof_FEC.Data[8286] := 619.71;
   Prof_FEC.Data[8287] := 685.0;
   Prof_FEC.Data[8288] := 617.21;
   Prof_FEC.Data[8289] := 604.94;
   Prof_FEC.Data[8290] := 701.15;
   Prof_FEC.Data[8291] := 642.22;
   Prof_FEC.Data[8292] := 591.7;
   Prof_FEC.Data[8293] := 567.72;
   Prof_FEC.Data[8294] := 570.38;
   Prof_FEC.Data[8295] := 573.09;
   Prof_FEC.Data[8296] := 652.99;
   Prof_FEC.Data[8297] := 576.33;
   Prof_FEC.Data[8298] := 542.96;
   Prof_FEC.Data[8299] := 591.89;
   Prof_FEC.Data[8300] := 501.74;
   Prof_FEC.Data[8301] := 474.6;
   Prof_FEC.Data[8302] := 490.15;
   Prof_FEC.Data[8303] := 587.71;
   Prof_FEC.Data[8304] := 567.01;
   Prof_FEC.Data[8305] := 617.85;
   Prof_FEC.Data[8306] := 632.44;
   Prof_FEC.Data[8307] := 649.22;
   Prof_FEC.Data[8308] := 645.48;
   Prof_FEC.Data[8309] := 596.12;
   Prof_FEC.Data[8310] := 581.23;
   Prof_FEC.Data[8311] := 552.59;
   Prof_FEC.Data[8312] := 550.69;
   Prof_FEC.Data[8313] := 641.74;
   Prof_FEC.Data[8314] := 582.68;
   Prof_FEC.Data[8315] := 535.44;
   Prof_FEC.Data[8316] := 625.92;
   Prof_FEC.Data[8317] := 612.53;
   Prof_FEC.Data[8318] := 616.47;
   Prof_FEC.Data[8319] := 457.76;
   Prof_FEC.Data[8320] := 282.93;
   Prof_FEC.Data[8321] := 204.65;
   Prof_FEC.Data[8322] := 153.26;
   Prof_FEC.Data[8323] := 126.49;
   Prof_FEC.Data[8324] := 107.79;
   Prof_FEC.Data[8325] := 87.64;
   Prof_FEC.Data[8326] := 91.39;
   Prof_FEC.Data[8327] := 108.77;
   Prof_FEC.Data[8328] := 183.75;
   Prof_FEC.Data[8329] := 192.21;
   Prof_FEC.Data[8330] := 193.92;
   Prof_FEC.Data[8331] := 204.61;
   Prof_FEC.Data[8332] := 38.275;
   Prof_FEC.Data[8333] := 38.408;
   Prof_FEC.Data[8334] := 37.717;
   Prof_FEC.Data[8335] := 41.171;
   Prof_FEC.Data[8336] := 40.373;
   Prof_FEC.Data[8337] := 39.781;
   Prof_FEC.Data[8338] := 39.567;
   Prof_FEC.Data[8339] := 40.069;
   Prof_FEC.Data[8340] := 40.536;
   Prof_FEC.Data[8341] := 39.149;
   Prof_FEC.Data[8342] := 38.345;
   Prof_FEC.Data[8343] := 38.813;
   Prof_FEC.Data[8344] := 38.705;
   Prof_FEC.Data[8345] := 35.505;
   Prof_FEC.Data[8346] := 39.912;
   Prof_FEC.Data[8347] := 39.485;
   Prof_FEC.Data[8348] := 40.9;
   Prof_FEC.Data[8349] := 39.103;
   Prof_FEC.Data[8350] := 40.085;
   Prof_FEC.Data[8351] := 40.846;
   Prof_FEC.Data[8352] := 41.325;
   Prof_FEC.Data[8353] := 41.463;
   Prof_FEC.Data[8354] := 41.976;
   Prof_FEC.Data[8355] := 39.423;
   Prof_FEC.Data[8356] := 40.153;
   Prof_FEC.Data[8357] := 40.75;
   Prof_FEC.Data[8358] := 40.928;
   Prof_FEC.Data[8359] := 39.712;
   Prof_FEC.Data[8360] := 46.289;
   Prof_FEC.Data[8361] := 44.657;
   Prof_FEC.Data[8362] := 46.856;
   Prof_FEC.Data[8363] := 45.304;
   Prof_FEC.Data[8364] := 43.516;
   Prof_FEC.Data[8365] := 42.853;
   Prof_FEC.Data[8366] := 40.608;
   Prof_FEC.Data[8367] := 40.579;
   Prof_FEC.Data[8368] := 42.405;
   Prof_FEC.Data[8369] := 42.285;
   Prof_FEC.Data[8370] := 45.782;
   Prof_FEC.Data[8371] := 42.906;
   Prof_FEC.Data[8372] := 264.28;
   Prof_FEC.Data[8373] := 234.03;
   Prof_FEC.Data[8374] := 263.07;
   Prof_FEC.Data[8375] := 249.77;
   Prof_FEC.Data[8376] := 311.34;
   Prof_FEC.Data[8377] := 278.75;
   Prof_FEC.Data[8378] := 306.99;
   Prof_FEC.Data[8379] := 299.65;
   Prof_FEC.Data[8380] := 290.77;
   Prof_FEC.Data[8381] := 307.35;
   Prof_FEC.Data[8382] := 318.1;
   Prof_FEC.Data[8383] := 328.72;
   Prof_FEC.Data[8384] := 342.47;
   Prof_FEC.Data[8385] := 406.67;
   Prof_FEC.Data[8386] := 415.35;
   Prof_FEC.Data[8387] := 406.6;
   Prof_FEC.Data[8388] := 396.82;
   Prof_FEC.Data[8389] := 371.17;
   Prof_FEC.Data[8390] := 356.54;
   Prof_FEC.Data[8391] := 335.03;
   Prof_FEC.Data[8392] := 339.04;
   Prof_FEC.Data[8393] := 357.59;
   Prof_FEC.Data[8394] := 304.13;
   Prof_FEC.Data[8395] := 323.43;
   Prof_FEC.Data[8396] := 284.43;
   Prof_FEC.Data[8397] := 245.11;
   Prof_FEC.Data[8398] := 249.71;
   Prof_FEC.Data[8399] := 244.96;
   Prof_FEC.Data[8400] := 270.75;
   Prof_FEC.Data[8401] := 248.76;
   Prof_FEC.Data[8402] := 259.01;
   Prof_FEC.Data[8403] := 279.79;
   Prof_FEC.Data[8404] := 302.24;
   Prof_FEC.Data[8405] := 295.58;
   Prof_FEC.Data[8406] := 286.27;
   Prof_FEC.Data[8407] := 287.35;
   Prof_FEC.Data[8408] := 309.08;
   Prof_FEC.Data[8409] := 301.6;
   Prof_FEC.Data[8410] := 298.14;
   Prof_FEC.Data[8411] := 237.24;
   Prof_FEC.Data[8412] := 149.84;
   Prof_FEC.Data[8413] := 122.17;
   Prof_FEC.Data[8414] := 110.98;
   Prof_FEC.Data[8415] := 102.24;
   Prof_FEC.Data[8416] := 122.42;
   Prof_FEC.Data[8417] := 111.27;
   Prof_FEC.Data[8418] := 117.36;
   Prof_FEC.Data[8419] := 120.42;
   Prof_FEC.Data[8420] := 117.48;
   Prof_FEC.Data[8421] := 117.58;
   Prof_FEC.Data[8422] := 114.85;
   Prof_FEC.Data[8423] := 161.89;
   Prof_FEC.Data[8424] := 176.72;
   Prof_FEC.Data[8425] := 186.37;
   Prof_FEC.Data[8426] := 234.88;
   Prof_FEC.Data[8427] := 208.19;
   Prof_FEC.Data[8428] := 38.382;
   Prof_FEC.Data[8429] := 39.604;
   Prof_FEC.Data[8430] := 40.466;
   Prof_FEC.Data[8431] := 39.914;
   Prof_FEC.Data[8432] := 39.113;
   Prof_FEC.Data[8433] := 39.577;
   Prof_FEC.Data[8434] := 37.77;
   Prof_FEC.Data[8435] := 41.621;
   Prof_FEC.Data[8436] := 41.028;
   Prof_FEC.Data[8437] := 40.265;
   Prof_FEC.Data[8438] := 41.435;
   Prof_FEC.Data[8439] := 42.024;
   Prof_FEC.Data[8440] := 38.954;
   Prof_FEC.Data[8441] := 40.418;
   Prof_FEC.Data[8442] := 41.998;
   Prof_FEC.Data[8443] := 43.337;
   Prof_FEC.Data[8444] := 44.831;
   Prof_FEC.Data[8445] := 43.412;
   Prof_FEC.Data[8446] := 43.701;
   Prof_FEC.Data[8447] := 42.549;
   Prof_FEC.Data[8448] := 42.817;
   Prof_FEC.Data[8449] := 41.163;
   Prof_FEC.Data[8450] := 41.949;
   Prof_FEC.Data[8451] := 39.213;
   Prof_FEC.Data[8452] := 41.971;
   Prof_FEC.Data[8453] := 46.371;
   Prof_FEC.Data[8454] := 44.733;
   Prof_FEC.Data[8455] := 46.428;
   Prof_FEC.Data[8456] := 42.433;
   Prof_FEC.Data[8457] := 41.829;
   Prof_FEC.Data[8458] := 44.583;
   Prof_FEC.Data[8459] := 44.25;
   Prof_FEC.Data[8460] := 46.64;
   Prof_FEC.Data[8461] := 46.106;
   Prof_FEC.Data[8462] := 46.719;
   Prof_FEC.Data[8463] := 50.0;
   Prof_FEC.Data[8464] := 45.821;
   Prof_FEC.Data[8465] := 44.873;
   Prof_FEC.Data[8466] := 44.613;
   Prof_FEC.Data[8467] := 45.332;
   Prof_FEC.Data[8468] := 293.83;
   Prof_FEC.Data[8469] := 355.24;
   Prof_FEC.Data[8470] := 321.05;
   Prof_FEC.Data[8471] := 270.59;
   Prof_FEC.Data[8472] := 187.22;
   Prof_FEC.Data[8473] := 155.45;
   Prof_FEC.Data[8474] := 145.48;
   Prof_FEC.Data[8475] := 168.0;
   Prof_FEC.Data[8476] := 196.69;
   Prof_FEC.Data[8477] := 218.19;
   Prof_FEC.Data[8478] := 194.67;
   Prof_FEC.Data[8479] := 179.41;
   Prof_FEC.Data[8480] := 156.66;
   Prof_FEC.Data[8481] := 150.69;
   Prof_FEC.Data[8482] := 142.91;
   Prof_FEC.Data[8483] := 150.15;
   Prof_FEC.Data[8484] := 172.47;
   Prof_FEC.Data[8485] := 186.24;
   Prof_FEC.Data[8486] := 176.0;
   Prof_FEC.Data[8487] := 168.64;
   Prof_FEC.Data[8488] := 146.74;
   Prof_FEC.Data[8489] := 145.64;
   Prof_FEC.Data[8490] := 135.4;
   Prof_FEC.Data[8491] := 141.52;
   Prof_FEC.Data[8492] := 142.97;
   Prof_FEC.Data[8493] := 147.61;
   Prof_FEC.Data[8494] := 121.76;
   Prof_FEC.Data[8495] := 148.93;
   Prof_FEC.Data[8496] := 116.05;
   Prof_FEC.Data[8497] := 111.35;
   Prof_FEC.Data[8498] := 109.75;
   Prof_FEC.Data[8499] := 115.92;
   Prof_FEC.Data[8500] := 134.12;
   Prof_FEC.Data[8501] := 142.28;
   Prof_FEC.Data[8502] := 139.34;
   Prof_FEC.Data[8503] := 143.06;
   Prof_FEC.Data[8504] := 118.39;
   Prof_FEC.Data[8505] := 115.86;
   Prof_FEC.Data[8506] := 120.08;
   Prof_FEC.Data[8507] := 112.32;
   Prof_FEC.Data[8508] := 131.79;
   Prof_FEC.Data[8509] := 134.4;
   Prof_FEC.Data[8510] := 143.29;
   Prof_FEC.Data[8511] := 130.19;
   Prof_FEC.Data[8512] := 139.18;
   Prof_FEC.Data[8513] := 126.09;
   Prof_FEC.Data[8514] := 126.34;
   Prof_FEC.Data[8515] := 115.84;
   Prof_FEC.Data[8516] := 121.46;
   Prof_FEC.Data[8517] := 122.13;
   Prof_FEC.Data[8518] := 138.74;
   Prof_FEC.Data[8519] := 158.41;
   Prof_FEC.Data[8520] := 181.88;
   Prof_FEC.Data[8521] := 194.92;
   Prof_FEC.Data[8522] := 205.32;
   Prof_FEC.Data[8523] := 266.35;
   Prof_FEC.Data[8524] := 42.232;
   Prof_FEC.Data[8525] := 43.903;
   Prof_FEC.Data[8526] := 43.44;
   Prof_FEC.Data[8527] := 46.294;
   Prof_FEC.Data[8528] := 43.498;
   Prof_FEC.Data[8529] := 40.584;
   Prof_FEC.Data[8530] := 42.796;
   Prof_FEC.Data[8531] := 42.641;
   Prof_FEC.Data[8532] := 42.483;
   Prof_FEC.Data[8533] := 47.089;
   Prof_FEC.Data[8534] := 46.219;
   Prof_FEC.Data[8535] := 44.223;
   Prof_FEC.Data[8536] := 44.544;
   Prof_FEC.Data[8537] := 44.876;
   Prof_FEC.Data[8538] := 42.509;
   Prof_FEC.Data[8539] := 44.226;
   Prof_FEC.Data[8540] := 46.103;
   Prof_FEC.Data[8541] := 44.863;
   Prof_FEC.Data[8542] := 44.372;
   Prof_FEC.Data[8543] := 44.147;
   Prof_FEC.Data[8544] := 43.204;
   Prof_FEC.Data[8545] := 43.269;
   Prof_FEC.Data[8546] := 39.222;
   Prof_FEC.Data[8547] := 40.191;
   Prof_FEC.Data[8548] := 44.433;
   Prof_FEC.Data[8549] := 46.729;
   Prof_FEC.Data[8550] := 47.42;
   Prof_FEC.Data[8551] := 45.957;
   Prof_FEC.Data[8552] := 43.177;
   Prof_FEC.Data[8553] := 42.281;
   Prof_FEC.Data[8554] := 41.821;
   Prof_FEC.Data[8555] := 43.703;
   Prof_FEC.Data[8556] := 41.606;
   Prof_FEC.Data[8557] := 45.476;
   Prof_FEC.Data[8558] := 46.197;
   Prof_FEC.Data[8559] := 42.113;
   Prof_FEC.Data[8560] := 41.585;
   Prof_FEC.Data[8561] := 40.895;
   Prof_FEC.Data[8562] := 41.3;
   Prof_FEC.Data[8563] := 42.044;
   Prof_FEC.Data[8564] := 382.92;
   Prof_FEC.Data[8565] := 378.9;
   Prof_FEC.Data[8566] := 407.86;
   Prof_FEC.Data[8567] := 343.36;
   Prof_FEC.Data[8568] := 387.67;
   Prof_FEC.Data[8569] := 360.8;
   Prof_FEC.Data[8570] := 464.66;
   Prof_FEC.Data[8571] := 428.57;
   Prof_FEC.Data[8572] := 560.98;
   Prof_FEC.Data[8573] := 588.02;
   Prof_FEC.Data[8574] := 607.19;
   Prof_FEC.Data[8575] := 688.74;
   Prof_FEC.Data[8576] := 656.09;
   Prof_FEC.Data[8577] := 667.94;
   Prof_FEC.Data[8578] := 755.12;
   Prof_FEC.Data[8579] := 675.22;
   Prof_FEC.Data[8580] := 652.23;
   Prof_FEC.Data[8581] := 655.5;
   Prof_FEC.Data[8582] := 615.07;
   Prof_FEC.Data[8583] := 707.42;
   Prof_FEC.Data[8584] := 686.18;
   Prof_FEC.Data[8585] := 606.21;
   Prof_FEC.Data[8586] := 600.05;
   Prof_FEC.Data[8587] := 617.79;
   Prof_FEC.Data[8588] := 643.5;
   Prof_FEC.Data[8589] := 598.43;
   Prof_FEC.Data[8590] := 540.79;
   Prof_FEC.Data[8591] := 540.43;
   Prof_FEC.Data[8592] := 584.37;
   Prof_FEC.Data[8593] := 647.96;
   Prof_FEC.Data[8594] := 629.3;
   Prof_FEC.Data[8595] := 676.58;
   Prof_FEC.Data[8596] := 668.51;
   Prof_FEC.Data[8597] := 638.76;
   Prof_FEC.Data[8598] := 623.16;
   Prof_FEC.Data[8599] := 573.31;
   Prof_FEC.Data[8600] := 582.97;
   Prof_FEC.Data[8601] := 547.12;
   Prof_FEC.Data[8602] := 617.2;
   Prof_FEC.Data[8603] := 585.91;
   Prof_FEC.Data[8604] := 653.92;
   Prof_FEC.Data[8605] := 636.43;
   Prof_FEC.Data[8606] := 595.36;
   Prof_FEC.Data[8607] := 474.1;
   Prof_FEC.Data[8608] := 321.96;
   Prof_FEC.Data[8609] := 209.88;
   Prof_FEC.Data[8610] := 161.98;
   Prof_FEC.Data[8611] := 140.39;
   Prof_FEC.Data[8612] := 119.46;
   Prof_FEC.Data[8613] := 88.59;
   Prof_FEC.Data[8614] := 85.51;
   Prof_FEC.Data[8615] := 108.87;
   Prof_FEC.Data[8616] := 174.22;
   Prof_FEC.Data[8617] := 225.24;
   Prof_FEC.Data[8618] := 226.11;
   Prof_FEC.Data[8619] := 218.05;
   Prof_FEC.Data[8620] := 37.379;
   Prof_FEC.Data[8621] := 40.237;
   Prof_FEC.Data[8622] := 39.091;
   Prof_FEC.Data[8623] := 39.829;
   Prof_FEC.Data[8624] := 39.681;
   Prof_FEC.Data[8625] := 40.919;
   Prof_FEC.Data[8626] := 39.845;
   Prof_FEC.Data[8627] := 42.445;
   Prof_FEC.Data[8628] := 41.237;
   Prof_FEC.Data[8629] := 39.903;
   Prof_FEC.Data[8630] := 39.109;
   Prof_FEC.Data[8631] := 37.336;
   Prof_FEC.Data[8632] := 41.253;
   Prof_FEC.Data[8633] := 41.314;
   Prof_FEC.Data[8634] := 40.602;
   Prof_FEC.Data[8635] := 40.692;
   Prof_FEC.Data[8636] := 39.774;
   Prof_FEC.Data[8637] := 39.017;
   Prof_FEC.Data[8638] := 37.928;
   Prof_FEC.Data[8639] := 38.909;
   Prof_FEC.Data[8640] := 43.918;
   Prof_FEC.Data[8641] := 42.288;
   Prof_FEC.Data[8642] := 40.496;
   Prof_FEC.Data[8643] := 43.038;
   Prof_FEC.Data[8644] := 38.584;
   Prof_FEC.Data[8645] := 41.3;
   Prof_FEC.Data[8646] := 38.967;
   Prof_FEC.Data[8647] := 39.889;
   Prof_FEC.Data[8648] := 41.654;
   Prof_FEC.Data[8649] := 43.17;
   Prof_FEC.Data[8650] := 41.786;
   Prof_FEC.Data[8651] := 42.584;
   Prof_FEC.Data[8652] := 38.497;
   Prof_FEC.Data[8653] := 38.856;
   Prof_FEC.Data[8654] := 39.58;
   Prof_FEC.Data[8655] := 41.352;
   Prof_FEC.Data[8656] := 41.197;
   Prof_FEC.Data[8657] := 44.142;
   Prof_FEC.Data[8658] := 46.632;
   Prof_FEC.Data[8659] := 48.277;
   Prof_FEC.Data[8660] := 376.75;
   Prof_FEC.Data[8661] := 449.11;
   Prof_FEC.Data[8662] := 416.45;
   Prof_FEC.Data[8663] := 487.64;
   Prof_FEC.Data[8664] := 433.69;
   Prof_FEC.Data[8665] := 478.63;
   Prof_FEC.Data[8666] := 436.45;
   Prof_FEC.Data[8667] := 482.32;
   Prof_FEC.Data[8668] := 579.17;
   Prof_FEC.Data[8669] := 634.32;
   Prof_FEC.Data[8670] := 606.56;
   Prof_FEC.Data[8671] := 648.9;
   Prof_FEC.Data[8672] := 697.16;
   Prof_FEC.Data[8673] := 729.01;
   Prof_FEC.Data[8674] := 688.12;
   Prof_FEC.Data[8675] := 709.76;
   Prof_FEC.Data[8676] := 660.06;
   Prof_FEC.Data[8677] := 713.2;
   Prof_FEC.Data[8678] := 740.23;
   Prof_FEC.Data[8679] := 695.98;
   Prof_FEC.Data[8680] := 662.31;
   Prof_FEC.Data[8681] := 744.24;
   Prof_FEC.Data[8682] := 597.49;
   Prof_FEC.Data[8683] := 673.27;
   Prof_FEC.Data[8684] := 645.06;
   Prof_FEC.Data[8685] := 627.61;
   Prof_FEC.Data[8686] := 598.55;
   Prof_FEC.Data[8687] := 631.67;
   Prof_FEC.Data[8688] := 641.22;
   Prof_FEC.Data[8689] := 649.4;
   Prof_FEC.Data[8690] := 569.18;
   Prof_FEC.Data[8691] := 698.35;
   Prof_FEC.Data[8692] := 649.48;
   Prof_FEC.Data[8693] := 631.31;
   Prof_FEC.Data[8694] := 608.62;
   Prof_FEC.Data[8695] := 665.94;
   Prof_FEC.Data[8696] := 609.3;
   Prof_FEC.Data[8697] := 586.9;
   Prof_FEC.Data[8698] := 635.96;
   Prof_FEC.Data[8699] := 635.82;
   Prof_FEC.Data[8700] := 658.38;
   Prof_FEC.Data[8701] := 680.11;
   Prof_FEC.Data[8702] := 640.08;
   Prof_FEC.Data[8703] := 494.1;
   Prof_FEC.Data[8704] := 303.35;
   Prof_FEC.Data[8705] := 204.0;
   Prof_FEC.Data[8706] := 133.78;
   Prof_FEC.Data[8707] := 119.18;
   Prof_FEC.Data[8708] := 91.73;
   Prof_FEC.Data[8709] := 74.04;
   Prof_FEC.Data[8710] := 69.58;
   Prof_FEC.Data[8711] := 86.4;
   Prof_FEC.Data[8712] := 142.83;
   Prof_FEC.Data[8713] := 180.22;
   Prof_FEC.Data[8714] := 185.36;
   Prof_FEC.Data[8715] := 198.59;
   Prof_FEC.Data[8716] := 37.143;
   Prof_FEC.Data[8717] := 40.451;
   Prof_FEC.Data[8718] := 40.749;
   Prof_FEC.Data[8719] := 40.145;
   Prof_FEC.Data[8720] := 42.058;
   Prof_FEC.Data[8721] := 40.255;
   Prof_FEC.Data[8722] := 39.887;
   Prof_FEC.Data[8723] := 42.045;
   Prof_FEC.Data[8724] := 40.306;
   Prof_FEC.Data[8725] := 40.685;
   Prof_FEC.Data[8726] := 37.99;
   Prof_FEC.Data[8727] := 37.369;
   Prof_FEC.Data[8728] := 38.643;
   Prof_FEC.Data[8729] := 36.372;
   Prof_FEC.Data[8730] := 37.39;
   Prof_FEC.Data[8731] := 38.238;
   Prof_FEC.Data[8732] := 36.38;
   Prof_FEC.Data[8733] := 32.6;
   Prof_FEC.Data[8734] := 33.635;
   Prof_FEC.Data[8735] := 35.016;
   Prof_FEC.Data[8736] := 37.082;
   Prof_FEC.Data[8737] := 36.614;
   Prof_FEC.Data[8738] := 35.677;
   Prof_FEC.Data[8739] := 34.776;
   Prof_FEC.Data[8740] := 32.581;
   Prof_FEC.Data[8741] := 33.275;
   Prof_FEC.Data[8742] := 35.534;
   Prof_FEC.Data[8743] := 34.845;
   Prof_FEC.Data[8744] := 36.631;
   Prof_FEC.Data[8745] := 35.309;
   Prof_FEC.Data[8746] := 37.643;
   Prof_FEC.Data[8747] := 37.241;
   Prof_FEC.Data[8748] := 36.162;
   Prof_FEC.Data[8749] := 37.128;
   Prof_FEC.Data[8750] := 37.884;
   Prof_FEC.Data[8751] := 35.153;
   Prof_FEC.Data[8752] := 36.377;
   Prof_FEC.Data[8753] := 36.242;
   Prof_FEC.Data[8754] := 37.226;
   Prof_FEC.Data[8755] := 41.834;
   Prof_FEC.Data[8756] := 329.23;
   Prof_FEC.Data[8757] := 420.06;
   Prof_FEC.Data[8758] := 360.67;
   Prof_FEC.Data[8759] := 471.2;
   Prof_FEC.Data[8760] := 369.87;
   Prof_FEC.Data[8761] := 396.88;
   Prof_FEC.Data[8762] := 397.98;
   Prof_FEC.Data[8763] := 511.31;
   Prof_FEC.Data[8764] := 490.33;
   Prof_FEC.Data[8765] := 513.24;
   Prof_FEC.Data[8766] := 615.27;
   Prof_FEC.Data[8767] := 610.72;
   Prof_FEC.Data[8768] := 598.77;
   Prof_FEC.Data[8769] := 605.67;
   Prof_FEC.Data[8770] := 615.61;
   Prof_FEC.Data[8771] := 727.3;
   Prof_FEC.Data[8772] := 694.85;
   Prof_FEC.Data[8773] := 711.12;
   Prof_FEC.Data[8774] := 709.57;
   Prof_FEC.Data[8775] := 612.0;
   Prof_FEC.Data[8776] := 664.14;
   Prof_FEC.Data[8777] := 639.75;
   Prof_FEC.Data[8778] := 685.7;
   Prof_FEC.Data[8779] := 587.11;
   Prof_FEC.Data[8780] := 624.04;
   Prof_FEC.Data[8781] := 644.81;
   Prof_FEC.Data[8782] := 519.18;
   Prof_FEC.Data[8783] := 598.6;
   Prof_FEC.Data[8784] := 634.04;
   Prof_FEC.Data[8785] := 682.97;
   Prof_FEC.Data[8786] := 581.28;
   Prof_FEC.Data[8787] := 676.23;
   Prof_FEC.Data[8788] := 654.85;
   Prof_FEC.Data[8789] := 666.78;
   Prof_FEC.Data[8790] := 743.03;
   Prof_FEC.Data[8791] := 632.97;
   Prof_FEC.Data[8792] := 675.69;
   Prof_FEC.Data[8793] := 654.39;
   Prof_FEC.Data[8794] := 681.35;
   Prof_FEC.Data[8795] := 703.44;
   Prof_FEC.Data[8796] := 764.34;
   Prof_FEC.Data[8797] := 682.82;
   Prof_FEC.Data[8798] := 665.13;
   Prof_FEC.Data[8799] := 529.25;
   Prof_FEC.Data[8800] := 273.92;
   Prof_FEC.Data[8801] := 189.9;
   Prof_FEC.Data[8802] := 150.29;
   Prof_FEC.Data[8803] := 119.93;
   Prof_FEC.Data[8804] := 105.31;
   Prof_FEC.Data[8805] := 74.48;
   Prof_FEC.Data[8806] := 71.7;
   Prof_FEC.Data[8807] := 98.06;
   Prof_FEC.Data[8808] := 158.69;
   Prof_FEC.Data[8809] := 183.1;
   Prof_FEC.Data[8810] := 185.55;
   Prof_FEC.Data[8811] := 213.32;
   Prof_FEC.Data[8812] := 38.51;
   Prof_FEC.Data[8813] := 38.039;
   Prof_FEC.Data[8814] := 37.207;
   Prof_FEC.Data[8815] := 38.178;
   Prof_FEC.Data[8816] := 40.716;
   Prof_FEC.Data[8817] := 39.019;
   Prof_FEC.Data[8818] := 40.537;
   Prof_FEC.Data[8819] := 39.172;
   Prof_FEC.Data[8820] := 38.074;
   Prof_FEC.Data[8821] := 39.524;
   Prof_FEC.Data[8822] := 37.604;
   Prof_FEC.Data[8823] := 37.889;
   Prof_FEC.Data[8824] := 38.892;
   Prof_FEC.Data[8825] := 39.286;
   Prof_FEC.Data[8826] := 41.291;
   Prof_FEC.Data[8827] := 40.539;
   Prof_FEC.Data[8828] := 39.752;
   Prof_FEC.Data[8829] := 38.567;
   Prof_FEC.Data[8830] := 38.156;
   Prof_FEC.Data[8831] := 39.491;
   Prof_FEC.Data[8832] := 39.425;
   Prof_FEC.Data[8833] := 41.999;
   Prof_FEC.Data[8834] := 41.205;
   Prof_FEC.Data[8835] := 39.472;
   Prof_FEC.Data[8836] := 37.846;
   Prof_FEC.Data[8837] := 39.172;
   Prof_FEC.Data[8838] := 39.1;
   Prof_FEC.Data[8839] := 38.285;
   Prof_FEC.Data[8840] := 39.74;
   Prof_FEC.Data[8841] := 40.599;
   Prof_FEC.Data[8842] := 39.205;
   Prof_FEC.Data[8843] := 40.136;
   Prof_FEC.Data[8844] := 37.292;
   Prof_FEC.Data[8845] := 36.336;
   Prof_FEC.Data[8846] := 37.363;
   Prof_FEC.Data[8847] := 36.107;
   Prof_FEC.Data[8848] := 35.235;
   Prof_FEC.Data[8849] := 37.554;
   Prof_FEC.Data[8850] := 39.551;
   Prof_FEC.Data[8851] := 40.684;
   Prof_FEC.Data[8852] := 302.43;
   Prof_FEC.Data[8853] := 392.33;
   Prof_FEC.Data[8854] := 402.62;
   Prof_FEC.Data[8855] := 406.09;
   Prof_FEC.Data[8856] := 386.24;
   Prof_FEC.Data[8857] := 448.69;
   Prof_FEC.Data[8858] := 427.39;
   Prof_FEC.Data[8859] := 433.68;
   Prof_FEC.Data[8860] := 568.39;
   Prof_FEC.Data[8861] := 566.55;
   Prof_FEC.Data[8862] := 622.09;
   Prof_FEC.Data[8863] := 656.75;
   Prof_FEC.Data[8864] := 639.66;
   Prof_FEC.Data[8865] := 627.21;
   Prof_FEC.Data[8866] := 690.53;
   Prof_FEC.Data[8867] := 738.29;
   Prof_FEC.Data[8868] := 691.64;
   Prof_FEC.Data[8869] := 679.74;
   Prof_FEC.Data[8870] := 707.03;
   Prof_FEC.Data[8871] := 641.21;
   Prof_FEC.Data[8872] := 643.7;
   Prof_FEC.Data[8873] := 628.12;
   Prof_FEC.Data[8874] := 639.81;
   Prof_FEC.Data[8875] := 629.72;
   Prof_FEC.Data[8876] := 651.11;
   Prof_FEC.Data[8877] := 656.84;
   Prof_FEC.Data[8878] := 623.54;
   Prof_FEC.Data[8879] := 569.13;
   Prof_FEC.Data[8880] := 685.92;
   Prof_FEC.Data[8881] := 791.15;
   Prof_FEC.Data[8882] := 777.69;
   Prof_FEC.Data[8883] := 771.06;
   Prof_FEC.Data[8884] := 743.0;
   Prof_FEC.Data[8885] := 769.49;
   Prof_FEC.Data[8886] := 734.03;
   Prof_FEC.Data[8887] := 714.45;
   Prof_FEC.Data[8888] := 629.64;
   Prof_FEC.Data[8889] := 668.76;
   Prof_FEC.Data[8890] := 642.61;
   Prof_FEC.Data[8891] := 639.0;
   Prof_FEC.Data[8892] := 620.04;
   Prof_FEC.Data[8893] := 669.97;
   Prof_FEC.Data[8894] := 618.81;
   Prof_FEC.Data[8895] := 499.04;
   Prof_FEC.Data[8896] := 266.3;
   Prof_FEC.Data[8897] := 157.31;
   Prof_FEC.Data[8898] := 136.26;
   Prof_FEC.Data[8899] := 114.31;
   Prof_FEC.Data[8900] := 72.26;
   Prof_FEC.Data[8901] := 58.55;
   Prof_FEC.Data[8902] := 62.69;
   Prof_FEC.Data[8903] := 80.63;
   Prof_FEC.Data[8904] := 133.57;
   Prof_FEC.Data[8905] := 152.05;
   Prof_FEC.Data[8906] := 145.44;
   Prof_FEC.Data[8907] := 161.51;
   Prof_FEC.Data[8908] := 34.055;
   Prof_FEC.Data[8909] := 34.027;
   Prof_FEC.Data[8910] := 35.086;
   Prof_FEC.Data[8911] := 36.6;
   Prof_FEC.Data[8912] := 36.519;
   Prof_FEC.Data[8913] := 37.416;
   Prof_FEC.Data[8914] := 36.93;
   Prof_FEC.Data[8915] := 37.53;
   Prof_FEC.Data[8916] := 37.445;
   Prof_FEC.Data[8917] := 37.241;
   Prof_FEC.Data[8918] := 37.887;
   Prof_FEC.Data[8919] := 36.949;
   Prof_FEC.Data[8920] := 40.221;
   Prof_FEC.Data[8921] := 41.459;
   Prof_FEC.Data[8922] := 40.254;
   Prof_FEC.Data[8923] := 40.629;
   Prof_FEC.Data[8924] := 40.91;
   Prof_FEC.Data[8925] := 37.885;
   Prof_FEC.Data[8926] := 37.434;
   Prof_FEC.Data[8927] := 40.303;
   Prof_FEC.Data[8928] := 41.561;
   Prof_FEC.Data[8929] := 41.556;
   Prof_FEC.Data[8930] := 40.179;
   Prof_FEC.Data[8931] := 40.486;
   Prof_FEC.Data[8932] := 38.075;
   Prof_FEC.Data[8933] := 40.107;
   Prof_FEC.Data[8934] := 40.986;
   Prof_FEC.Data[8935] := 41.195;
   Prof_FEC.Data[8936] := 41.565;
   Prof_FEC.Data[8937] := 41.969;
   Prof_FEC.Data[8938] := 44.119;
   Prof_FEC.Data[8939] := 38.773;
   Prof_FEC.Data[8940] := 39.095;
   Prof_FEC.Data[8941] := 38.007;
   Prof_FEC.Data[8942] := 40.352;
   Prof_FEC.Data[8943] := 38.316;
   Prof_FEC.Data[8944] := 39.928;
   Prof_FEC.Data[8945] := 39.544;
   Prof_FEC.Data[8946] := 42.169;
   Prof_FEC.Data[8947] := 45.319;
   Prof_FEC.Data[8948] := 362.66;
   Prof_FEC.Data[8949] := 398.42;
   Prof_FEC.Data[8950] := 438.08;
   Prof_FEC.Data[8951] := 429.88;
   Prof_FEC.Data[8952] := 425.74;
   Prof_FEC.Data[8953] := 432.17;
   Prof_FEC.Data[8954] := 409.0;
   Prof_FEC.Data[8955] := 501.7;
   Prof_FEC.Data[8956] := 493.53;
   Prof_FEC.Data[8957] := 478.69;
   Prof_FEC.Data[8958] := 503.76;
   Prof_FEC.Data[8959] := 550.43;
   Prof_FEC.Data[8960] := 529.95;
   Prof_FEC.Data[8961] := 545.26;
   Prof_FEC.Data[8962] := 476.56;
   Prof_FEC.Data[8963] := 598.19;
   Prof_FEC.Data[8964] := 607.45;
   Prof_FEC.Data[8965] := 564.53;
   Prof_FEC.Data[8966] := 597.15;
   Prof_FEC.Data[8967] := 590.35;
   Prof_FEC.Data[8968] := 567.83;
   Prof_FEC.Data[8969] := 545.62;
   Prof_FEC.Data[8970] := 590.19;
   Prof_FEC.Data[8971] := 613.1;
   Prof_FEC.Data[8972] := 619.18;
   Prof_FEC.Data[8973] := 468.31;
   Prof_FEC.Data[8974] := 523.91;
   Prof_FEC.Data[8975] := 477.41;
   Prof_FEC.Data[8976] := 558.72;
   Prof_FEC.Data[8977] := 563.55;
   Prof_FEC.Data[8978] := 654.56;
   Prof_FEC.Data[8979] := 562.29;
   Prof_FEC.Data[8980] := 614.98;
   Prof_FEC.Data[8981] := 630.04;
   Prof_FEC.Data[8982] := 598.12;
   Prof_FEC.Data[8983] := 606.01;
   Prof_FEC.Data[8984] := 614.02;
   Prof_FEC.Data[8985] := 609.42;
   Prof_FEC.Data[8986] := 596.49;
   Prof_FEC.Data[8987] := 610.89;
   Prof_FEC.Data[8988] := 672.06;
   Prof_FEC.Data[8989] := 670.03;
   Prof_FEC.Data[8990] := 659.19;
   Prof_FEC.Data[8991] := 517.99;
   Prof_FEC.Data[8992] := 293.28;
   Prof_FEC.Data[8993] := 188.77;
   Prof_FEC.Data[8994] := 141.68;
   Prof_FEC.Data[8995] := 125.9;
   Prof_FEC.Data[8996] := 97.59;
   Prof_FEC.Data[8997] := 71.44;
   Prof_FEC.Data[8998] := 70.29;
   Prof_FEC.Data[8999] := 91.41;
   Prof_FEC.Data[9000] := 155.62;
   Prof_FEC.Data[9001] := 175.29;
   Prof_FEC.Data[9002] := 190.24;
   Prof_FEC.Data[9003] := 192.4;
   Prof_FEC.Data[9004] := 37.473;
   Prof_FEC.Data[9005] := 37.167;
   Prof_FEC.Data[9006] := 39.277;
   Prof_FEC.Data[9007] := 40.154;
   Prof_FEC.Data[9008] := 39.985;
   Prof_FEC.Data[9009] := 40.096;
   Prof_FEC.Data[9010] := 39.478;
   Prof_FEC.Data[9011] := 38.156;
   Prof_FEC.Data[9012] := 37.981;
   Prof_FEC.Data[9013] := 36.899;
   Prof_FEC.Data[9014] := 37.649;
   Prof_FEC.Data[9015] := 41.273;
   Prof_FEC.Data[9016] := 40.777;
   Prof_FEC.Data[9017] := 42.382;
   Prof_FEC.Data[9018] := 39.209;
   Prof_FEC.Data[9019] := 39.893;
   Prof_FEC.Data[9020] := 39.67;
   Prof_FEC.Data[9021] := 39.263;
   Prof_FEC.Data[9022] := 38.054;
   Prof_FEC.Data[9023] := 40.067;
   Prof_FEC.Data[9024] := 42.334;
   Prof_FEC.Data[9025] := 42.359;
   Prof_FEC.Data[9026] := 43.028;
   Prof_FEC.Data[9027] := 42.528;
   Prof_FEC.Data[9028] := 40.926;
   Prof_FEC.Data[9029] := 38.264;
   Prof_FEC.Data[9030] := 37.212;
   Prof_FEC.Data[9031] := 39.502;
   Prof_FEC.Data[9032] := 42.935;
   Prof_FEC.Data[9033] := 41.991;
   Prof_FEC.Data[9034] := 40.324;
   Prof_FEC.Data[9035] := 42.937;
   Prof_FEC.Data[9036] := 41.091;
   Prof_FEC.Data[9037] := 36.331;
   Prof_FEC.Data[9038] := 38.876;
   Prof_FEC.Data[9039] := 38.468;
   Prof_FEC.Data[9040] := 38.039;
   Prof_FEC.Data[9041] := 38.604;
   Prof_FEC.Data[9042] := 39.55;
   Prof_FEC.Data[9043] := 37.93;
   Prof_FEC.Data[9044] := 205.37;
   Prof_FEC.Data[9045] := 198.17;
   Prof_FEC.Data[9046] := 215.35;
   Prof_FEC.Data[9047] := 222.81;
   Prof_FEC.Data[9048] := 243.57;
   Prof_FEC.Data[9049] := 253.02;
   Prof_FEC.Data[9050] := 253.96;
   Prof_FEC.Data[9051] := 257.96;
   Prof_FEC.Data[9052] := 280.49;
   Prof_FEC.Data[9053] := 279.62;
   Prof_FEC.Data[9054] := 271.83;
   Prof_FEC.Data[9055] := 284.89;
   Prof_FEC.Data[9056] := 353.97;
   Prof_FEC.Data[9057] := 362.75;
   Prof_FEC.Data[9058] := 389.09;
   Prof_FEC.Data[9059] := 391.12;
   Prof_FEC.Data[9060] := 351.9;
   Prof_FEC.Data[9061] := 350.35;
   Prof_FEC.Data[9062] := 316.07;
   Prof_FEC.Data[9063] := 336.99;
   Prof_FEC.Data[9064] := 373.95;
   Prof_FEC.Data[9065] := 320.71;
   Prof_FEC.Data[9066] := 373.11;
   Prof_FEC.Data[9067] := 324.88;
   Prof_FEC.Data[9068] := 345.85;
   Prof_FEC.Data[9069] := 314.89;
   Prof_FEC.Data[9070] := 290.4;
   Prof_FEC.Data[9071] := 262.7;
   Prof_FEC.Data[9072] := 284.91;
   Prof_FEC.Data[9073] := 291.8;
   Prof_FEC.Data[9074] := 244.15;
   Prof_FEC.Data[9075] := 276.99;
   Prof_FEC.Data[9076] := 282.88;
   Prof_FEC.Data[9077] := 250.6;
   Prof_FEC.Data[9078] := 285.78;
   Prof_FEC.Data[9079] := 282.57;
   Prof_FEC.Data[9080] := 334.35;
   Prof_FEC.Data[9081] := 301.03;
   Prof_FEC.Data[9082] := 292.03;
   Prof_FEC.Data[9083] := 229.07;
   Prof_FEC.Data[9084] := 104.05;
   Prof_FEC.Data[9085] := 81.03;
   Prof_FEC.Data[9086] := 65.58;
   Prof_FEC.Data[9087] := 59.25;
   Prof_FEC.Data[9088] := 82.69;
   Prof_FEC.Data[9089] := 78.16;
   Prof_FEC.Data[9090] := 78.81;
   Prof_FEC.Data[9091] := 86.35;
   Prof_FEC.Data[9092] := 81.28;
   Prof_FEC.Data[9093] := 84.92;
   Prof_FEC.Data[9094] := 92.52;
   Prof_FEC.Data[9095] := 98.7;
   Prof_FEC.Data[9096] := 106.83;
   Prof_FEC.Data[9097] := 131.78;
   Prof_FEC.Data[9098] := 143.98;
   Prof_FEC.Data[9099] := 176.5;
   Prof_FEC.Data[9100] := 34.828;
   Prof_FEC.Data[9101] := 37.017;
   Prof_FEC.Data[9102] := 38.899;
   Prof_FEC.Data[9103] := 41.491;
   Prof_FEC.Data[9104] := 37.646;
   Prof_FEC.Data[9105] := 40.249;
   Prof_FEC.Data[9106] := 40.75;
   Prof_FEC.Data[9107] := 38.428;
   Prof_FEC.Data[9108] := 40.058;
   Prof_FEC.Data[9109] := 41.705;
   Prof_FEC.Data[9110] := 43.421;
   Prof_FEC.Data[9111] := 39.978;
   Prof_FEC.Data[9112] := 40.976;
   Prof_FEC.Data[9113] := 39.57;
   Prof_FEC.Data[9114] := 38.273;
   Prof_FEC.Data[9115] := 38.517;
   Prof_FEC.Data[9116] := 41.41;
   Prof_FEC.Data[9117] := 43.471;
   Prof_FEC.Data[9118] := 40.41;
   Prof_FEC.Data[9119] := 40.078;
   Prof_FEC.Data[9120] := 38.522;
   Prof_FEC.Data[9121] := 40.073;
   Prof_FEC.Data[9122] := 38.634;
   Prof_FEC.Data[9123] := 39.706;
   Prof_FEC.Data[9124] := 44.184;
   Prof_FEC.Data[9125] := 41.726;
   Prof_FEC.Data[9126] := 38.503;
   Prof_FEC.Data[9127] := 39.802;
   Prof_FEC.Data[9128] := 38.814;
   Prof_FEC.Data[9129] := 36.602;
   Prof_FEC.Data[9130] := 36.879;
   Prof_FEC.Data[9131] := 36.792;
   Prof_FEC.Data[9132] := 37.97;
   Prof_FEC.Data[9133] := 37.625;
   Prof_FEC.Data[9134] := 36.233;
   Prof_FEC.Data[9135] := 35.952;
   Prof_FEC.Data[9136] := 38.857;
   Prof_FEC.Data[9137] := 37.757;
   Prof_FEC.Data[9138] := 38.636;
   Prof_FEC.Data[9139] := 35.992;
   Prof_FEC.Data[9140] := 218.83;
   Prof_FEC.Data[9141] := 239.86;
   Prof_FEC.Data[9142] := 225.22;
   Prof_FEC.Data[9143] := 186.8;
   Prof_FEC.Data[9144] := 136.19;
   Prof_FEC.Data[9145] := 116.82;
   Prof_FEC.Data[9146] := 98.98;
   Prof_FEC.Data[9147] := 104.36;
   Prof_FEC.Data[9148] := 130.01;
   Prof_FEC.Data[9149] := 131.32;
   Prof_FEC.Data[9150] := 136.19;
   Prof_FEC.Data[9151] := 122.82;
   Prof_FEC.Data[9152] := 108.61;
   Prof_FEC.Data[9153] := 112.11;
   Prof_FEC.Data[9154] := 99.37;
   Prof_FEC.Data[9155] := 117.3;
   Prof_FEC.Data[9156] := 118.54;
   Prof_FEC.Data[9157] := 132.28;
   Prof_FEC.Data[9158] := 113.24;
   Prof_FEC.Data[9159] := 113.4;
   Prof_FEC.Data[9160] := 96.04;
   Prof_FEC.Data[9161] := 88.29;
   Prof_FEC.Data[9162] := 93.31;
   Prof_FEC.Data[9163] := 91.52;
   Prof_FEC.Data[9164] := 94.08;
   Prof_FEC.Data[9165] := 94.26;
   Prof_FEC.Data[9166] := 93.36;
   Prof_FEC.Data[9167] := 95.08;
   Prof_FEC.Data[9168] := 69.03;
   Prof_FEC.Data[9169] := 70.01;
   Prof_FEC.Data[9170] := 83.82;
   Prof_FEC.Data[9171] := 89.75;
   Prof_FEC.Data[9172] := 83.65;
   Prof_FEC.Data[9173] := 80.49;
   Prof_FEC.Data[9174] := 89.36;
   Prof_FEC.Data[9175] := 80.7;
   Prof_FEC.Data[9176] := 78.02;
   Prof_FEC.Data[9177] := 78.05;
   Prof_FEC.Data[9178] := 73.41;
   Prof_FEC.Data[9179] := 86.57;
   Prof_FEC.Data[9180] := 92.95;
   Prof_FEC.Data[9181] := 94.0;
   Prof_FEC.Data[9182] := 95.27;
   Prof_FEC.Data[9183] := 100.99;
   Prof_FEC.Data[9184] := 89.31;
   Prof_FEC.Data[9185] := 92.67;
   Prof_FEC.Data[9186] := 90.15;
   Prof_FEC.Data[9187] := 85.11;
   Prof_FEC.Data[9188] := 100.18;
   Prof_FEC.Data[9189] := 109.53;
   Prof_FEC.Data[9190] := 119.76;
   Prof_FEC.Data[9191] := 112.81;
   Prof_FEC.Data[9192] := 121.76;
   Prof_FEC.Data[9193] := 162.05;
   Prof_FEC.Data[9194] := 167.52;
   Prof_FEC.Data[9195] := 190.76;
   Prof_FEC.Data[9196] := 39.759;
   Prof_FEC.Data[9197] := 41.651;
   Prof_FEC.Data[9198] := 42.855;
   Prof_FEC.Data[9199] := 43.531;
   Prof_FEC.Data[9200] := 42.321;
   Prof_FEC.Data[9201] := 40.717;
   Prof_FEC.Data[9202] := 40.699;
   Prof_FEC.Data[9203] := 40.336;
   Prof_FEC.Data[9204] := 39.54;
   Prof_FEC.Data[9205] := 42.303;
   Prof_FEC.Data[9206] := 42.442;
   Prof_FEC.Data[9207] := 41.18;
   Prof_FEC.Data[9208] := 39.947;
   Prof_FEC.Data[9209] := 38.8;
   Prof_FEC.Data[9210] := 39.556;
   Prof_FEC.Data[9211] := 42.017;
   Prof_FEC.Data[9212] := 42.881;
   Prof_FEC.Data[9213] := 43.808;
   Prof_FEC.Data[9214] := 38.817;
   Prof_FEC.Data[9215] := 39.285;
   Prof_FEC.Data[9216] := 39.237;
   Prof_FEC.Data[9217] := 40.884;
   Prof_FEC.Data[9218] := 37.478;
   Prof_FEC.Data[9219] := 38.273;
   Prof_FEC.Data[9220] := 38.337;
   Prof_FEC.Data[9221] := 40.608;
   Prof_FEC.Data[9222] := 38.41;
   Prof_FEC.Data[9223] := 39.886;
   Prof_FEC.Data[9224] := 35.495;
   Prof_FEC.Data[9225] := 34.189;
   Prof_FEC.Data[9226] := 40.045;
   Prof_FEC.Data[9227] := 37.842;
   Prof_FEC.Data[9228] := 43.563;
   Prof_FEC.Data[9229] := 44.542;
   Prof_FEC.Data[9230] := 40.237;
   Prof_FEC.Data[9231] := 40.591;
   Prof_FEC.Data[9232] := 36.734;
   Prof_FEC.Data[9233] := 38.901;
   Prof_FEC.Data[9234] := 39.015;
   Prof_FEC.Data[9235] := 42.293;
   Prof_FEC.Data[9236] := 321.9;
   Prof_FEC.Data[9237] := 350.48;
   Prof_FEC.Data[9238] := 407.72;
   Prof_FEC.Data[9239] := 379.81;
   Prof_FEC.Data[9240] := 383.55;
   Prof_FEC.Data[9241] := 430.03;
   Prof_FEC.Data[9242] := 430.01;
   Prof_FEC.Data[9243] := 439.21;
   Prof_FEC.Data[9244] := 528.46;
   Prof_FEC.Data[9245] := 522.87;
   Prof_FEC.Data[9246] := 612.72;
   Prof_FEC.Data[9247] := 547.04;
   Prof_FEC.Data[9248] := 698.12;
   Prof_FEC.Data[9249] := 693.9;
   Prof_FEC.Data[9250] := 726.11;
   Prof_FEC.Data[9251] := 743.05;
   Prof_FEC.Data[9252] := 696.52;
   Prof_FEC.Data[9253] := 657.02;
   Prof_FEC.Data[9254] := 679.63;
   Prof_FEC.Data[9255] := 793.93;
   Prof_FEC.Data[9256] := 701.04;
   Prof_FEC.Data[9257] := 669.31;
   Prof_FEC.Data[9258] := 711.0;
   Prof_FEC.Data[9259] := 668.8;
   Prof_FEC.Data[9260] := 621.82;
   Prof_FEC.Data[9261] := 566.2;
   Prof_FEC.Data[9262] := 607.61;
   Prof_FEC.Data[9263] := 611.78;
   Prof_FEC.Data[9264] := 613.44;
   Prof_FEC.Data[9265] := 618.4;
   Prof_FEC.Data[9266] := 577.86;
   Prof_FEC.Data[9267] := 657.11;
   Prof_FEC.Data[9268] := 626.51;
   Prof_FEC.Data[9269] := 643.29;
   Prof_FEC.Data[9270] := 716.52;
   Prof_FEC.Data[9271] := 632.61;
   Prof_FEC.Data[9272] := 640.75;
   Prof_FEC.Data[9273] := 730.73;
   Prof_FEC.Data[9274] := 623.07;
   Prof_FEC.Data[9275] := 678.03;
   Prof_FEC.Data[9276] := 681.03;
   Prof_FEC.Data[9277] := 706.8;
   Prof_FEC.Data[9278] := 749.58;
   Prof_FEC.Data[9279] := 565.05;
   Prof_FEC.Data[9280] := 339.26;
   Prof_FEC.Data[9281] := 246.51;
   Prof_FEC.Data[9282] := 165.56;
   Prof_FEC.Data[9283] := 147.14;
   Prof_FEC.Data[9284] := 118.35;
   Prof_FEC.Data[9285] := 89.85;
   Prof_FEC.Data[9286] := 76.83;
   Prof_FEC.Data[9287] := 99.32;
   Prof_FEC.Data[9288] := 153.25;
   Prof_FEC.Data[9289] := 184.29;
   Prof_FEC.Data[9290] := 194.04;
   Prof_FEC.Data[9291] := 221.48;
   Prof_FEC.Data[9292] := 37.282;
   Prof_FEC.Data[9293] := 36.993;
   Prof_FEC.Data[9294] := 38.433;
   Prof_FEC.Data[9295] := 38.099;
   Prof_FEC.Data[9296] := 36.932;
   Prof_FEC.Data[9297] := 39.516;
   Prof_FEC.Data[9298] := 39.705;
   Prof_FEC.Data[9299] := 41.626;
   Prof_FEC.Data[9300] := 38.186;
   Prof_FEC.Data[9301] := 38.594;
   Prof_FEC.Data[9302] := 38.057;
   Prof_FEC.Data[9303] := 40.195;
   Prof_FEC.Data[9304] := 37.824;
   Prof_FEC.Data[9305] := 40.454;
   Prof_FEC.Data[9306] := 41.313;
   Prof_FEC.Data[9307] := 39.316;
   Prof_FEC.Data[9308] := 41.554;
   Prof_FEC.Data[9309] := 37.606;
   Prof_FEC.Data[9310] := 38.491;
   Prof_FEC.Data[9311] := 40.108;
   Prof_FEC.Data[9312] := 38.447;
   Prof_FEC.Data[9313] := 38.722;
   Prof_FEC.Data[9314] := 38.651;
   Prof_FEC.Data[9315] := 37.412;
   Prof_FEC.Data[9316] := 36.77;
   Prof_FEC.Data[9317] := 34.592;
   Prof_FEC.Data[9318] := 33.303;
   Prof_FEC.Data[9319] := 36.823;
   Prof_FEC.Data[9320] := 36.617;
   Prof_FEC.Data[9321] := 37.896;
   Prof_FEC.Data[9322] := 38.295;
   Prof_FEC.Data[9323] := 36.375;
   Prof_FEC.Data[9324] := 34.562;
   Prof_FEC.Data[9325] := 36.309;
   Prof_FEC.Data[9326] := 35.26;
   Prof_FEC.Data[9327] := 37.177;
   Prof_FEC.Data[9328] := 33.975;
   Prof_FEC.Data[9329] := 35.914;
   Prof_FEC.Data[9330] := 35.381;
   Prof_FEC.Data[9331] := 40.828;
   Prof_FEC.Data[9332] := 272.05;
   Prof_FEC.Data[9333] := 350.79;
   Prof_FEC.Data[9334] := 393.0;
   Prof_FEC.Data[9335] := 421.35;
   Prof_FEC.Data[9336] := 351.55;
   Prof_FEC.Data[9337] := 384.16;
   Prof_FEC.Data[9338] := 460.37;
   Prof_FEC.Data[9339] := 445.97;
   Prof_FEC.Data[9340] := 468.64;
   Prof_FEC.Data[9341] := 527.81;
   Prof_FEC.Data[9342] := 534.35;
   Prof_FEC.Data[9343] := 525.45;
   Prof_FEC.Data[9344] := 583.12;
   Prof_FEC.Data[9345] := 551.87;
   Prof_FEC.Data[9346] := 608.0;
   Prof_FEC.Data[9347] := 573.36;
   Prof_FEC.Data[9348] := 628.39;
   Prof_FEC.Data[9349] := 728.45;
   Prof_FEC.Data[9350] := 612.21;
   Prof_FEC.Data[9351] := 651.55;
   Prof_FEC.Data[9352] := 659.58;
   Prof_FEC.Data[9353] := 647.65;
   Prof_FEC.Data[9354] := 625.26;
   Prof_FEC.Data[9355] := 641.22;
   Prof_FEC.Data[9356] := 590.53;
   Prof_FEC.Data[9357] := 560.94;
   Prof_FEC.Data[9358] := 481.51;
   Prof_FEC.Data[9359] := 573.83;
   Prof_FEC.Data[9360] := 586.45;
   Prof_FEC.Data[9361] := 592.9;
   Prof_FEC.Data[9362] := 566.97;
   Prof_FEC.Data[9363] := 578.72;
   Prof_FEC.Data[9364] := 605.3;
   Prof_FEC.Data[9365] := 630.87;
   Prof_FEC.Data[9366] := 589.51;
   Prof_FEC.Data[9367] := 580.03;
   Prof_FEC.Data[9368] := 586.0;
   Prof_FEC.Data[9369] := 604.88;
   Prof_FEC.Data[9370] := 596.68;
   Prof_FEC.Data[9371] := 537.34;
   Prof_FEC.Data[9372] := 592.0;
   Prof_FEC.Data[9373] := 604.14;
   Prof_FEC.Data[9374] := 608.8;
   Prof_FEC.Data[9375] := 398.85;
   Prof_FEC.Data[9376] := 191.85;
   Prof_FEC.Data[9377] := 145.72;
   Prof_FEC.Data[9378] := 80.18;
   Prof_FEC.Data[9379] := 81.28;
   Prof_FEC.Data[9380] := 47.11;
   Prof_FEC.Data[9381] := 35.49;
   Prof_FEC.Data[9382] := 32.34;
   Prof_FEC.Data[9383] := 43.91;
   Prof_FEC.Data[9384] := 84.89;
   Prof_FEC.Data[9385] := 82.89;
   Prof_FEC.Data[9386] := 96.85;
   Prof_FEC.Data[9387] := 114.7;
   Prof_FEC.Data[9388] := 31.194;
   Prof_FEC.Data[9389] := 33.341;
   Prof_FEC.Data[9390] := 34.447;
   Prof_FEC.Data[9391] := 34.332;
   Prof_FEC.Data[9392] := 31.285;
   Prof_FEC.Data[9393] := 31.643;
   Prof_FEC.Data[9394] := 32.301;
   Prof_FEC.Data[9395] := 33.463;
   Prof_FEC.Data[9396] := 33.017;
   Prof_FEC.Data[9397] := 31.726;
   Prof_FEC.Data[9398] := 33.726;
   Prof_FEC.Data[9399] := 34.502;
   Prof_FEC.Data[9400] := 33.056;
   Prof_FEC.Data[9401] := 33.171;
   Prof_FEC.Data[9402] := 33.515;
   Prof_FEC.Data[9403] := 34.077;
   Prof_FEC.Data[9404] := 35.076;
   Prof_FEC.Data[9405] := 34.569;
   Prof_FEC.Data[9406] := 38.115;
   Prof_FEC.Data[9407] := 35.496;
   Prof_FEC.Data[9408] := 37.717;
   Prof_FEC.Data[9409] := 35.305;
   Prof_FEC.Data[9410] := 38.35;
   Prof_FEC.Data[9411] := 37.67;
   Prof_FEC.Data[9412] := 37.244;
   Prof_FEC.Data[9413] := 35.282;
   Prof_FEC.Data[9414] := 37.779;
   Prof_FEC.Data[9415] := 37.871;
   Prof_FEC.Data[9416] := 40.196;
   Prof_FEC.Data[9417] := 38.938;
   Prof_FEC.Data[9418] := 41.021;
   Prof_FEC.Data[9419] := 41.228;
   Prof_FEC.Data[9420] := 39.376;
   Prof_FEC.Data[9421] := 41.421;
   Prof_FEC.Data[9422] := 39.854;
   Prof_FEC.Data[9423] := 39.179;
   Prof_FEC.Data[9424] := 38.724;
   Prof_FEC.Data[9425] := 40.506;
   Prof_FEC.Data[9426] := 39.751;
   Prof_FEC.Data[9427] := 40.105;
   Prof_FEC.Data[9428] := 310.91;
   Prof_FEC.Data[9429] := 370.02;
   Prof_FEC.Data[9430] := 424.31;
   Prof_FEC.Data[9431] := 466.78;
   Prof_FEC.Data[9432] := 473.89;
   Prof_FEC.Data[9433] := 467.74;
   Prof_FEC.Data[9434] := 496.73;
   Prof_FEC.Data[9435] := 519.68;
   Prof_FEC.Data[9436] := 515.67;
   Prof_FEC.Data[9437] := 597.95;
   Prof_FEC.Data[9438] := 576.03;
   Prof_FEC.Data[9439] := 644.92;
   Prof_FEC.Data[9440] := 683.17;
   Prof_FEC.Data[9441] := 700.06;
   Prof_FEC.Data[9442] := 710.5;
   Prof_FEC.Data[9443] := 719.01;
   Prof_FEC.Data[9444] := 758.49;
   Prof_FEC.Data[9445] := 734.47;
   Prof_FEC.Data[9446] := 741.38;
   Prof_FEC.Data[9447] := 792.75;
   Prof_FEC.Data[9448] := 796.7;
   Prof_FEC.Data[9449] := 746.47;
   Prof_FEC.Data[9450] := 734.71;
   Prof_FEC.Data[9451] := 744.97;
   Prof_FEC.Data[9452] := 697.24;
   Prof_FEC.Data[9453] := 641.63;
   Prof_FEC.Data[9454] := 606.8;
   Prof_FEC.Data[9455] := 650.08;
   Prof_FEC.Data[9456] := 680.73;
   Prof_FEC.Data[9457] := 724.14;
   Prof_FEC.Data[9458] := 722.26;
   Prof_FEC.Data[9459] := 673.78;
   Prof_FEC.Data[9460] := 647.07;
   Prof_FEC.Data[9461] := 661.42;
   Prof_FEC.Data[9462] := 580.95;
   Prof_FEC.Data[9463] := 597.26;
   Prof_FEC.Data[9464] := 594.93;
   Prof_FEC.Data[9465] := 625.34;
   Prof_FEC.Data[9466] := 576.46;
   Prof_FEC.Data[9467] := 613.26;
   Prof_FEC.Data[9468] := 674.32;
   Prof_FEC.Data[9469] := 715.63;
   Prof_FEC.Data[9470] := 624.68;
   Prof_FEC.Data[9471] := 460.34;
   Prof_FEC.Data[9472] := 249.84;
   Prof_FEC.Data[9473] := 177.85;
   Prof_FEC.Data[9474] := 124.69;
   Prof_FEC.Data[9475] := 108.17;
   Prof_FEC.Data[9476] := 89.72;
   Prof_FEC.Data[9477] := 72.69;
   Prof_FEC.Data[9478] := 68.28;
   Prof_FEC.Data[9479] := 78.71;
   Prof_FEC.Data[9480] := 118.99;
   Prof_FEC.Data[9481] := 153.52;
   Prof_FEC.Data[9482] := 144.92;
   Prof_FEC.Data[9483] := 162.42;
   Prof_FEC.Data[9484] := 33.969;
   Prof_FEC.Data[9485] := 37.115;
   Prof_FEC.Data[9486] := 35.726;
   Prof_FEC.Data[9487] := 35.841;
   Prof_FEC.Data[9488] := 36.399;
   Prof_FEC.Data[9489] := 37.419;
   Prof_FEC.Data[9490] := 39.146;
   Prof_FEC.Data[9491] := 36.174;
   Prof_FEC.Data[9492] := 35.081;
   Prof_FEC.Data[9493] := 34.6;
   Prof_FEC.Data[9494] := 35.773;
   Prof_FEC.Data[9495] := 40.074;
   Prof_FEC.Data[9496] := 39.605;
   Prof_FEC.Data[9497] := 40.244;
   Prof_FEC.Data[9498] := 40.387;
   Prof_FEC.Data[9499] := 39.543;
   Prof_FEC.Data[9500] := 38.248;
   Prof_FEC.Data[9501] := 35.579;
   Prof_FEC.Data[9502] := 35.58;
   Prof_FEC.Data[9503] := 35.203;
   Prof_FEC.Data[9504] := 36.276;
   Prof_FEC.Data[9505] := 36.3;
   Prof_FEC.Data[9506] := 35.759;
   Prof_FEC.Data[9507] := 38.57;
   Prof_FEC.Data[9508] := 35.873;
   Prof_FEC.Data[9509] := 34.252;
   Prof_FEC.Data[9510] := 33.587;
   Prof_FEC.Data[9511] := 34.998;
   Prof_FEC.Data[9512] := 35.822;
   Prof_FEC.Data[9513] := 37.82;
   Prof_FEC.Data[9514] := 37.427;
   Prof_FEC.Data[9515] := 37.389;
   Prof_FEC.Data[9516] := 36.255;
   Prof_FEC.Data[9517] := 37.068;
   Prof_FEC.Data[9518] := 36.098;
   Prof_FEC.Data[9519] := 35.701;
   Prof_FEC.Data[9520] := 37.655;
   Prof_FEC.Data[9521] := 37.197;
   Prof_FEC.Data[9522] := 36.872;
   Prof_FEC.Data[9523] := 37.383;
   Prof_FEC.Data[9524] := 257.5;
   Prof_FEC.Data[9525] := 293.92;
   Prof_FEC.Data[9526] := 344.0;
   Prof_FEC.Data[9527] := 367.3;
   Prof_FEC.Data[9528] := 357.48;
   Prof_FEC.Data[9529] := 423.92;
   Prof_FEC.Data[9530] := 429.69;
   Prof_FEC.Data[9531] := 441.46;
   Prof_FEC.Data[9532] := 511.39;
   Prof_FEC.Data[9533] := 546.75;
   Prof_FEC.Data[9534] := 565.06;
   Prof_FEC.Data[9535] := 572.08;
   Prof_FEC.Data[9536] := 578.84;
   Prof_FEC.Data[9537] := 561.76;
   Prof_FEC.Data[9538] := 610.95;
   Prof_FEC.Data[9539] := 704.33;
   Prof_FEC.Data[9540] := 611.07;
   Prof_FEC.Data[9541] := 613.54;
   Prof_FEC.Data[9542] := 689.78;
   Prof_FEC.Data[9543] := 694.39;
   Prof_FEC.Data[9544] := 684.89;
   Prof_FEC.Data[9545] := 691.66;
   Prof_FEC.Data[9546] := 743.29;
   Prof_FEC.Data[9547] := 739.52;
   Prof_FEC.Data[9548] := 672.28;
   Prof_FEC.Data[9549] := 697.93;
   Prof_FEC.Data[9550] := 689.19;
   Prof_FEC.Data[9551] := 637.07;
   Prof_FEC.Data[9552] := 749.62;
   Prof_FEC.Data[9553] := 762.54;
   Prof_FEC.Data[9554] := 664.04;
   Prof_FEC.Data[9555] := 751.65;
   Prof_FEC.Data[9556] := 658.08;
   Prof_FEC.Data[9557] := 661.87;
   Prof_FEC.Data[9558] := 753.79;
   Prof_FEC.Data[9559] := 764.77;
   Prof_FEC.Data[9560] := 726.84;
   Prof_FEC.Data[9561] := 722.51;
   Prof_FEC.Data[9562] := 720.46;
   Prof_FEC.Data[9563] := 731.58;
   Prof_FEC.Data[9564] := 798.16;
   Prof_FEC.Data[9565] := 739.18;
   Prof_FEC.Data[9566] := 687.11;
   Prof_FEC.Data[9567] := 560.0;
   Prof_FEC.Data[9568] := 331.54;
   Prof_FEC.Data[9569] := 230.65;
   Prof_FEC.Data[9570] := 164.14;
   Prof_FEC.Data[9571] := 133.62;
   Prof_FEC.Data[9572] := 123.86;
   Prof_FEC.Data[9573] := 93.27;
   Prof_FEC.Data[9574] := 86.87;
   Prof_FEC.Data[9575] := 110.63;
   Prof_FEC.Data[9576] := 148.75;
   Prof_FEC.Data[9577] := 170.7;
   Prof_FEC.Data[9578] := 171.53;
   Prof_FEC.Data[9579] := 190.6;
   Prof_FEC.Data[9580] := 34.452;
   Prof_FEC.Data[9581] := 35.536;
   Prof_FEC.Data[9582] := 37.109;
   Prof_FEC.Data[9583] := 36.498;
   Prof_FEC.Data[9584] := 38.428;
   Prof_FEC.Data[9585] := 37.028;
   Prof_FEC.Data[9586] := 37.289;
   Prof_FEC.Data[9587] := 39.157;
   Prof_FEC.Data[9588] := 39.462;
   Prof_FEC.Data[9589] := 35.756;
   Prof_FEC.Data[9590] := 36.861;
   Prof_FEC.Data[9591] := 36.708;
   Prof_FEC.Data[9592] := 36.232;
   Prof_FEC.Data[9593] := 38.245;
   Prof_FEC.Data[9594] := 36.337;
   Prof_FEC.Data[9595] := 36.435;
   Prof_FEC.Data[9596] := 36.716;
   Prof_FEC.Data[9597] := 37.985;
   Prof_FEC.Data[9598] := 35.752;
   Prof_FEC.Data[9599] := 39.808;
   Prof_FEC.Data[9600] := 38.062;
   Prof_FEC.Data[9601] := 40.696;
   Prof_FEC.Data[9602] := 40.079;
   Prof_FEC.Data[9603] := 40.499;
   Prof_FEC.Data[9604] := 40.55;
   Prof_FEC.Data[9605] := 37.651;
   Prof_FEC.Data[9606] := 38.245;
   Prof_FEC.Data[9607] := 37.647;
   Prof_FEC.Data[9608] := 38.697;
   Prof_FEC.Data[9609] := 38.551;
   Prof_FEC.Data[9610] := 38.656;
   Prof_FEC.Data[9611] := 36.931;
   Prof_FEC.Data[9612] := 35.252;
   Prof_FEC.Data[9613] := 32.116;
   Prof_FEC.Data[9614] := 38.006;
   Prof_FEC.Data[9615] := 39.107;
   Prof_FEC.Data[9616] := 39.66;
   Prof_FEC.Data[9617] := 36.706;
   Prof_FEC.Data[9618] := 38.013;
   Prof_FEC.Data[9619] := 39.797;
   Prof_FEC.Data[9620] := 324.89;
   Prof_FEC.Data[9621] := 370.45;
   Prof_FEC.Data[9622] := 371.08;
   Prof_FEC.Data[9623] := 405.13;
   Prof_FEC.Data[9624] := 393.66;
   Prof_FEC.Data[9625] := 394.63;
   Prof_FEC.Data[9626] := 432.99;
   Prof_FEC.Data[9627] := 479.54;
   Prof_FEC.Data[9628] := 481.48;
   Prof_FEC.Data[9629] := 557.78;
   Prof_FEC.Data[9630] := 555.55;
   Prof_FEC.Data[9631] := 571.29;
   Prof_FEC.Data[9632] := 642.97;
   Prof_FEC.Data[9633] := 730.36;
   Prof_FEC.Data[9634] := 779.14;
   Prof_FEC.Data[9635] := 700.61;
   Prof_FEC.Data[9636] := 739.47;
   Prof_FEC.Data[9637] := 689.32;
   Prof_FEC.Data[9638] := 694.9;
   Prof_FEC.Data[9639] := 666.97;
   Prof_FEC.Data[9640] := 705.75;
   Prof_FEC.Data[9641] := 689.01;
   Prof_FEC.Data[9642] := 638.41;
   Prof_FEC.Data[9643] := 666.2;
   Prof_FEC.Data[9644] := 591.55;
   Prof_FEC.Data[9645] := 580.13;
   Prof_FEC.Data[9646] := 564.87;
   Prof_FEC.Data[9647] := 597.24;
   Prof_FEC.Data[9648] := 650.22;
   Prof_FEC.Data[9649] := 649.82;
   Prof_FEC.Data[9650] := 629.4;
   Prof_FEC.Data[9651] := 587.46;
   Prof_FEC.Data[9652] := 570.06;
   Prof_FEC.Data[9653] := 548.22;
   Prof_FEC.Data[9654] := 585.89;
   Prof_FEC.Data[9655] := 571.48;
   Prof_FEC.Data[9656] := 658.16;
   Prof_FEC.Data[9657] := 650.96;
   Prof_FEC.Data[9658] := 642.93;
   Prof_FEC.Data[9659] := 583.8;
   Prof_FEC.Data[9660] := 680.69;
   Prof_FEC.Data[9661] := 624.64;
   Prof_FEC.Data[9662] := 635.03;
   Prof_FEC.Data[9663] := 482.21;
   Prof_FEC.Data[9664] := 222.95;
   Prof_FEC.Data[9665] := 154.43;
   Prof_FEC.Data[9666] := 97.93;
   Prof_FEC.Data[9667] := 83.72;
   Prof_FEC.Data[9668] := 67.37;
   Prof_FEC.Data[9669] := 53.66;
   Prof_FEC.Data[9670] := 51.62;
   Prof_FEC.Data[9671] := 59.15;
   Prof_FEC.Data[9672] := 98.56;
   Prof_FEC.Data[9673] := 96.26;
   Prof_FEC.Data[9674] := 140.99;
   Prof_FEC.Data[9675] := 139.91;
   Prof_FEC.Data[9676] := 31.03;
   Prof_FEC.Data[9677] := 33.528;
   Prof_FEC.Data[9678] := 30.602;
   Prof_FEC.Data[9679] := 32.578;
   Prof_FEC.Data[9680] := 33.332;
   Prof_FEC.Data[9681] := 35.131;
   Prof_FEC.Data[9682] := 33.692;
   Prof_FEC.Data[9683] := 35.261;
   Prof_FEC.Data[9684] := 33.155;
   Prof_FEC.Data[9685] := 33.485;
   Prof_FEC.Data[9686] := 33.811;
   Prof_FEC.Data[9687] := 33.681;
   Prof_FEC.Data[9688] := 34.546;
   Prof_FEC.Data[9689] := 33.771;
   Prof_FEC.Data[9690] := 34.44;
   Prof_FEC.Data[9691] := 33.26;
   Prof_FEC.Data[9692] := 33.298;
   Prof_FEC.Data[9693] := 33.951;
   Prof_FEC.Data[9694] := 33.52;
   Prof_FEC.Data[9695] := 33.36;
   Prof_FEC.Data[9696] := 31.719;
   Prof_FEC.Data[9697] := 34.018;
   Prof_FEC.Data[9698] := 34.363;
   Prof_FEC.Data[9699] := 35.062;
   Prof_FEC.Data[9700] := 34.985;
   Prof_FEC.Data[9701] := 32.842;
   Prof_FEC.Data[9702] := 33.534;
   Prof_FEC.Data[9703] := 33.693;
   Prof_FEC.Data[9704] := 33.707;
   Prof_FEC.Data[9705] := 33.677;
   Prof_FEC.Data[9706] := 30.854;
   Prof_FEC.Data[9707] := 32.386;
   Prof_FEC.Data[9708] := 34.967;
   Prof_FEC.Data[9709] := 34.953;
   Prof_FEC.Data[9710] := 35.99;
   Prof_FEC.Data[9711] := 36.546;
   Prof_FEC.Data[9712] := 37.081;
   Prof_FEC.Data[9713] := 35.747;
   Prof_FEC.Data[9714] := 36.319;
   Prof_FEC.Data[9715] := 35.891;
   Prof_FEC.Data[9716] := 145.67;
   Prof_FEC.Data[9717] := 124.11;
   Prof_FEC.Data[9718] := 140.59;
   Prof_FEC.Data[9719] := 163.09;
   Prof_FEC.Data[9720] := 197.82;
   Prof_FEC.Data[9721] := 229.15;
   Prof_FEC.Data[9722] := 248.26;
   Prof_FEC.Data[9723] := 262.83;
   Prof_FEC.Data[9724] := 262.1;
   Prof_FEC.Data[9725] := 253.73;
   Prof_FEC.Data[9726] := 238.04;
   Prof_FEC.Data[9727] := 324.73;
   Prof_FEC.Data[9728] := 294.62;
   Prof_FEC.Data[9729] := 283.03;
   Prof_FEC.Data[9730] := 296.93;
   Prof_FEC.Data[9731] := 301.13;
   Prof_FEC.Data[9732] := 288.35;
   Prof_FEC.Data[9733] := 318.27;
   Prof_FEC.Data[9734] := 283.14;
   Prof_FEC.Data[9735] := 354.98;
   Prof_FEC.Data[9736] := 359.8;
   Prof_FEC.Data[9737] := 339.94;
   Prof_FEC.Data[9738] := 344.48;
   Prof_FEC.Data[9739] := 287.59;
   Prof_FEC.Data[9740] := 254.41;
   Prof_FEC.Data[9741] := 247.28;
   Prof_FEC.Data[9742] := 233.96;
   Prof_FEC.Data[9743] := 226.44;
   Prof_FEC.Data[9744] := 241.41;
   Prof_FEC.Data[9745] := 258.53;
   Prof_FEC.Data[9746] := 285.97;
   Prof_FEC.Data[9747] := 269.01;
   Prof_FEC.Data[9748] := 241.42;
   Prof_FEC.Data[9749] := 241.85;
   Prof_FEC.Data[9750] := 232.53;
   Prof_FEC.Data[9751] := 274.05;
   Prof_FEC.Data[9752] := 295.82;
   Prof_FEC.Data[9753] := 324.63;
   Prof_FEC.Data[9754] := 261.97;
   Prof_FEC.Data[9755] := 201.62;
   Prof_FEC.Data[9756] := 93.22;
   Prof_FEC.Data[9757] := 54.51;
   Prof_FEC.Data[9758] := 40.62;
   Prof_FEC.Data[9759] := 42.52;
   Prof_FEC.Data[9760] := 64.57;
   Prof_FEC.Data[9761] := 60.56;
   Prof_FEC.Data[9762] := 68.14;
   Prof_FEC.Data[9763] := 65.31;
   Prof_FEC.Data[9764] := 65.35;
   Prof_FEC.Data[9765] := 66.4;
   Prof_FEC.Data[9766] := 72.7;
   Prof_FEC.Data[9767] := 91.38;
   Prof_FEC.Data[9768] := 95.18;
   Prof_FEC.Data[9769] := 114.84;
   Prof_FEC.Data[9770] := 132.11;
   Prof_FEC.Data[9771] := 153.74;
   Prof_FEC.Data[9772] := 33.382;
   Prof_FEC.Data[9773] := 36.09;
   Prof_FEC.Data[9774] := 36.612;
   Prof_FEC.Data[9775] := 36.594;
   Prof_FEC.Data[9776] := 37.723;
   Prof_FEC.Data[9777] := 35.745;
   Prof_FEC.Data[9778] := 34.982;
   Prof_FEC.Data[9779] := 37.379;
   Prof_FEC.Data[9780] := 37.56;
   Prof_FEC.Data[9781] := 36.817;
   Prof_FEC.Data[9782] := 36.277;
   Prof_FEC.Data[9783] := 37.486;
   Prof_FEC.Data[9784] := 35.405;
   Prof_FEC.Data[9785] := 37.019;
   Prof_FEC.Data[9786] := 34.966;
   Prof_FEC.Data[9787] := 36.712;
   Prof_FEC.Data[9788] := 36.326;
   Prof_FEC.Data[9789] := 35.711;
   Prof_FEC.Data[9790] := 32.853;
   Prof_FEC.Data[9791] := 33.248;
   Prof_FEC.Data[9792] := 36.291;
   Prof_FEC.Data[9793] := 34.835;
   Prof_FEC.Data[9794] := 33.26;
   Prof_FEC.Data[9795] := 33.852;
   Prof_FEC.Data[9796] := 33.8;
   Prof_FEC.Data[9797] := 32.361;
   Prof_FEC.Data[9798] := 34.71;
   Prof_FEC.Data[9799] := 34.205;
   Prof_FEC.Data[9800] := 32.8;
   Prof_FEC.Data[9801] := 33.475;
   Prof_FEC.Data[9802] := 34.1;
   Prof_FEC.Data[9803] := 34.646;
   Prof_FEC.Data[9804] := 34.625;
   Prof_FEC.Data[9805] := 34.414;
   Prof_FEC.Data[9806] := 33.505;
   Prof_FEC.Data[9807] := 36.095;
   Prof_FEC.Data[9808] := 34.932;
   Prof_FEC.Data[9809] := 37.844;
   Prof_FEC.Data[9810] := 36.534;
   Prof_FEC.Data[9811] := 32.676;
   Prof_FEC.Data[9812] := 148.55;
   Prof_FEC.Data[9813] := 129.54;
   Prof_FEC.Data[9814] := 118.24;
   Prof_FEC.Data[9815] := 104.71;
   Prof_FEC.Data[9816] := 81.28;
   Prof_FEC.Data[9817] := 64.93;
   Prof_FEC.Data[9818] := 69.27;
   Prof_FEC.Data[9819] := 59.63;
   Prof_FEC.Data[9820] := 66.47;
   Prof_FEC.Data[9821] := 62.43;
   Prof_FEC.Data[9822] := 64.77;
   Prof_FEC.Data[9823] := 68.19;
   Prof_FEC.Data[9824] := 71.72;
   Prof_FEC.Data[9825] := 64.07;
   Prof_FEC.Data[9826] := 58.92;
   Prof_FEC.Data[9827] := 63.47;
   Prof_FEC.Data[9828] := 62.88;
   Prof_FEC.Data[9829] := 63.09;
   Prof_FEC.Data[9830] := 64.66;
   Prof_FEC.Data[9831] := 62.0;
   Prof_FEC.Data[9832] := 69.29;
   Prof_FEC.Data[9833] := 59.8;
   Prof_FEC.Data[9834] := 66.14;
   Prof_FEC.Data[9835] := 63.99;
   Prof_FEC.Data[9836] := 69.05;
   Prof_FEC.Data[9837] := 69.59;
   Prof_FEC.Data[9838] := 73.54;
   Prof_FEC.Data[9839] := 79.63;
   Prof_FEC.Data[9840] := 76.15;
   Prof_FEC.Data[9841] := 80.11;
   Prof_FEC.Data[9842] := 82.12;
   Prof_FEC.Data[9843] := 90.95;
   Prof_FEC.Data[9844] := 85.4;
   Prof_FEC.Data[9845] := 85.54;
   Prof_FEC.Data[9846] := 81.69;
   Prof_FEC.Data[9847] := 98.1;
   Prof_FEC.Data[9848] := 94.04;
   Prof_FEC.Data[9849] := 100.5;
   Prof_FEC.Data[9850] := 89.02;
   Prof_FEC.Data[9851] := 93.04;
   Prof_FEC.Data[9852] := 85.25;
   Prof_FEC.Data[9853] := 88.75;
   Prof_FEC.Data[9854] := 89.75;
   Prof_FEC.Data[9855] := 88.95;
   Prof_FEC.Data[9856] := 85.87;
   Prof_FEC.Data[9857] := 89.0;
   Prof_FEC.Data[9858] := 89.57;
   Prof_FEC.Data[9859] := 93.66;
   Prof_FEC.Data[9860] := 82.5;
   Prof_FEC.Data[9861] := 84.36;
   Prof_FEC.Data[9862] := 91.7;
   Prof_FEC.Data[9863] := 109.89;
   Prof_FEC.Data[9864] := 131.05;
   Prof_FEC.Data[9865] := 133.47;
   Prof_FEC.Data[9866] := 149.52;
   Prof_FEC.Data[9867] := 170.67;
   Prof_FEC.Data[9868] := 34.958;
   Prof_FEC.Data[9869] := 39.645;
   Prof_FEC.Data[9870] := 38.72;
   Prof_FEC.Data[9871] := 37.993;
   Prof_FEC.Data[9872] := 38.113;
   Prof_FEC.Data[9873] := 37.763;
   Prof_FEC.Data[9874] := 36.025;
   Prof_FEC.Data[9875] := 37.509;
   Prof_FEC.Data[9876] := 38.464;
   Prof_FEC.Data[9877] := 38.053;
   Prof_FEC.Data[9878] := 35.255;
   Prof_FEC.Data[9879] := 37.177;
   Prof_FEC.Data[9880] := 36.599;
   Prof_FEC.Data[9881] := 39.215;
   Prof_FEC.Data[9882] := 39.252;
   Prof_FEC.Data[9883] := 38.407;
   Prof_FEC.Data[9884] := 36.586;
   Prof_FEC.Data[9885] := 38.803;
   Prof_FEC.Data[9886] := 35.641;
   Prof_FEC.Data[9887] := 39.199;
   Prof_FEC.Data[9888] := 37.711;
   Prof_FEC.Data[9889] := 38.481;
   Prof_FEC.Data[9890] := 39.459;
   Prof_FEC.Data[9891] := 37.357;
   Prof_FEC.Data[9892] := 39.537;
   Prof_FEC.Data[9893] := 39.438;
   Prof_FEC.Data[9894] := 39.211;
   Prof_FEC.Data[9895] := 38.261;
   Prof_FEC.Data[9896] := 43.008;
   Prof_FEC.Data[9897] := 40.455;
   Prof_FEC.Data[9898] := 40.065;
   Prof_FEC.Data[9899] := 39.04;
   Prof_FEC.Data[9900] := 37.462;
   Prof_FEC.Data[9901] := 39.96;
   Prof_FEC.Data[9902] := 38.793;
   Prof_FEC.Data[9903] := 37.092;
   Prof_FEC.Data[9904] := 37.079;
   Prof_FEC.Data[9905] := 36.394;
   Prof_FEC.Data[9906] := 39.308;
   Prof_FEC.Data[9907] := 40.819;
   Prof_FEC.Data[9908] := 284.36;
   Prof_FEC.Data[9909] := 336.1;
   Prof_FEC.Data[9910] := 354.03;
   Prof_FEC.Data[9911] := 392.86;
   Prof_FEC.Data[9912] := 412.72;
   Prof_FEC.Data[9913] := 395.83;
   Prof_FEC.Data[9914] := 437.82;
   Prof_FEC.Data[9915] := 404.56;
   Prof_FEC.Data[9916] := 487.82;
   Prof_FEC.Data[9917] := 481.98;
   Prof_FEC.Data[9918] := 526.82;
   Prof_FEC.Data[9919] := 545.45;
   Prof_FEC.Data[9920] := 568.56;
   Prof_FEC.Data[9921] := 605.54;
   Prof_FEC.Data[9922] := 725.4;
   Prof_FEC.Data[9923] := 694.62;
   Prof_FEC.Data[9924] := 608.13;
   Prof_FEC.Data[9925] := 665.49;
   Prof_FEC.Data[9926] := 630.13;
   Prof_FEC.Data[9927] := 668.87;
   Prof_FEC.Data[9928] := 647.12;
   Prof_FEC.Data[9929] := 693.53;
   Prof_FEC.Data[9930] := 702.69;
   Prof_FEC.Data[9931] := 652.56;
   Prof_FEC.Data[9932] := 615.54;
   Prof_FEC.Data[9933] := 588.4;
   Prof_FEC.Data[9934] := 556.87;
   Prof_FEC.Data[9935] := 576.75;
   Prof_FEC.Data[9936] := 667.21;
   Prof_FEC.Data[9937] := 715.45;
   Prof_FEC.Data[9938] := 611.8;
   Prof_FEC.Data[9939] := 693.04;
   Prof_FEC.Data[9940] := 659.94;
   Prof_FEC.Data[9941] := 702.47;
   Prof_FEC.Data[9942] := 648.84;
   Prof_FEC.Data[9943] := 587.16;
   Prof_FEC.Data[9944] := 648.66;
   Prof_FEC.Data[9945] := 602.75;
   Prof_FEC.Data[9946] := 626.74;
   Prof_FEC.Data[9947] := 620.3;
   Prof_FEC.Data[9948] := 680.27;
   Prof_FEC.Data[9949] := 655.86;
   Prof_FEC.Data[9950] := 559.43;
   Prof_FEC.Data[9951] := 484.29;
   Prof_FEC.Data[9952] := 265.37;
   Prof_FEC.Data[9953] := 178.5;
   Prof_FEC.Data[9954] := 130.65;
   Prof_FEC.Data[9955] := 111.91;
   Prof_FEC.Data[9956] := 87.17;
   Prof_FEC.Data[9957] := 69.35;
   Prof_FEC.Data[9958] := 66.92;
   Prof_FEC.Data[9959] := 85.38;
   Prof_FEC.Data[9960] := 113.89;
   Prof_FEC.Data[9961] := 147.76;
   Prof_FEC.Data[9962] := 155.91;
   Prof_FEC.Data[9963] := 192.84;
   Prof_FEC.Data[9964] := 36.626;
   Prof_FEC.Data[9965] := 37.397;
   Prof_FEC.Data[9966] := 40.005;
   Prof_FEC.Data[9967] := 40.256;
   Prof_FEC.Data[9968] := 40.604;
   Prof_FEC.Data[9969] := 38.132;
   Prof_FEC.Data[9970] := 39.921;
   Prof_FEC.Data[9971] := 39.683;
   Prof_FEC.Data[9972] := 39.897;
   Prof_FEC.Data[9973] := 38.607;
   Prof_FEC.Data[9974] := 38.117;
   Prof_FEC.Data[9975] := 37.843;
   Prof_FEC.Data[9976] := 40.683;
   Prof_FEC.Data[9977] := 41.553;
   Prof_FEC.Data[9978] := 39.004;
   Prof_FEC.Data[9979] := 39.477;
   Prof_FEC.Data[9980] := 37.921;
   Prof_FEC.Data[9981] := 36.635;
   Prof_FEC.Data[9982] := 39.601;
   Prof_FEC.Data[9983] := 38.622;
   Prof_FEC.Data[9984] := 39.791;
   Prof_FEC.Data[9985] := 42.644;
   Prof_FEC.Data[9986] := 39.281;
   Prof_FEC.Data[9987] := 38.479;
   Prof_FEC.Data[9988] := 39.144;
   Prof_FEC.Data[9989] := 38.068;
   Prof_FEC.Data[9990] := 40.541;
   Prof_FEC.Data[9991] := 42.998;
   Prof_FEC.Data[9992] := 45.185;
   Prof_FEC.Data[9993] := 46.224;
   Prof_FEC.Data[9994] := 44.081;
   Prof_FEC.Data[9995] := 42.988;
   Prof_FEC.Data[9996] := 41.834;
   Prof_FEC.Data[9997] := 43.43;
   Prof_FEC.Data[9998] := 41.791;
   Prof_FEC.Data[9999] := 41.407;
   Prof_FEC.Data[10000] := 45.805;
   Prof_FEC.Data[10001] := 45.866;
   Prof_FEC.Data[10002] := 47.467;
   Prof_FEC.Data[10003] := 48.597;
   Prof_FEC.Data[10004] := 354.3;
   Prof_FEC.Data[10005] := 366.44;
   Prof_FEC.Data[10006] := 378.76;
   Prof_FEC.Data[10007] := 415.22;
   Prof_FEC.Data[10008] := 454.74;
   Prof_FEC.Data[10009] := 479.05;
   Prof_FEC.Data[10010] := 479.83;
   Prof_FEC.Data[10011] := 498.99;
   Prof_FEC.Data[10012] := 541.5;
   Prof_FEC.Data[10013] := 666.0;
   Prof_FEC.Data[10014] := 704.44;
   Prof_FEC.Data[10015] := 727.89;
   Prof_FEC.Data[10016] := 761.59;
   Prof_FEC.Data[10017] := 776.05;
   Prof_FEC.Data[10018] := 758.38;
   Prof_FEC.Data[10019] := 755.82;
   Prof_FEC.Data[10020] := 697.96;
   Prof_FEC.Data[10021] := 701.89;
   Prof_FEC.Data[10022] := 715.68;
   Prof_FEC.Data[10023] := 716.33;
   Prof_FEC.Data[10024] := 707.82;
   Prof_FEC.Data[10025] := 709.11;
   Prof_FEC.Data[10026] := 645.69;
   Prof_FEC.Data[10027] := 617.6;
   Prof_FEC.Data[10028] := 634.32;
   Prof_FEC.Data[10029] := 601.18;
   Prof_FEC.Data[10030] := 599.01;
   Prof_FEC.Data[10031] := 625.11;
   Prof_FEC.Data[10032] := 643.45;
   Prof_FEC.Data[10033] := 570.52;
   Prof_FEC.Data[10034] := 649.67;
   Prof_FEC.Data[10035] := 704.25;
   Prof_FEC.Data[10036] := 727.16;
   Prof_FEC.Data[10037] := 788.83;
   Prof_FEC.Data[10038] := 729.21;
   Prof_FEC.Data[10039] := 681.44;
   Prof_FEC.Data[10040] := 676.8;
   Prof_FEC.Data[10041] := 680.21;
   Prof_FEC.Data[10042] := 664.24;
   Prof_FEC.Data[10043] := 716.12;
   Prof_FEC.Data[10044] := 813.34;
   Prof_FEC.Data[10045] := 780.21;
   Prof_FEC.Data[10046] := 668.28;
   Prof_FEC.Data[10047] := 542.26;
   Prof_FEC.Data[10048] := 280.72;
   Prof_FEC.Data[10049] := 210.18;
   Prof_FEC.Data[10050] := 147.79;
   Prof_FEC.Data[10051] := 110.76;
   Prof_FEC.Data[10052] := 100.24;
   Prof_FEC.Data[10053] := 76.56;
   Prof_FEC.Data[10054] := 71.52;
   Prof_FEC.Data[10055] := 78.14;
   Prof_FEC.Data[10056] := 103.05;
   Prof_FEC.Data[10057] := 143.35;
   Prof_FEC.Data[10058] := 156.78;
   Prof_FEC.Data[10059] := 170.32;
   Prof_FEC.Data[10060] := 36.124;
   Prof_FEC.Data[10061] := 37.499;
   Prof_FEC.Data[10062] := 38.371;
   Prof_FEC.Data[10063] := 37.883;
   Prof_FEC.Data[10064] := 37.091;
   Prof_FEC.Data[10065] := 38.848;
   Prof_FEC.Data[10066] := 39.304;
   Prof_FEC.Data[10067] := 38.334;
   Prof_FEC.Data[10068] := 38.039;
   Prof_FEC.Data[10069] := 36.494;
   Prof_FEC.Data[10070] := 37.217;
   Prof_FEC.Data[10071] := 36.896;
   Prof_FEC.Data[10072] := 38.932;
   Prof_FEC.Data[10073] := 38.786;
   Prof_FEC.Data[10074] := 37.675;
   Prof_FEC.Data[10075] := 39.975;
   Prof_FEC.Data[10076] := 40.239;
   Prof_FEC.Data[10077] := 38.792;
   Prof_FEC.Data[10078] := 38.243;
   Prof_FEC.Data[10079] := 38.219;
   Prof_FEC.Data[10080] := 39.531;
   Prof_FEC.Data[10081] := 41.382;
   Prof_FEC.Data[10082] := 42.321;
   Prof_FEC.Data[10083] := 42.236;
   Prof_FEC.Data[10084] := 39.901;
   Prof_FEC.Data[10085] := 39.847;
   Prof_FEC.Data[10086] := 40.278;
   Prof_FEC.Data[10087] := 40.373;
   Prof_FEC.Data[10088] := 42.464;
   Prof_FEC.Data[10089] := 41.261;
   Prof_FEC.Data[10090] := 41.533;
   Prof_FEC.Data[10091] := 40.038;
   Prof_FEC.Data[10092] := 38.877;
   Prof_FEC.Data[10093] := 37.781;
   Prof_FEC.Data[10094] := 35.623;
   Prof_FEC.Data[10095] := 38.564;
   Prof_FEC.Data[10096] := 37.847;
   Prof_FEC.Data[10097] := 36.456;
   Prof_FEC.Data[10098] := 38.698;
   Prof_FEC.Data[10099] := 42.525;
   Prof_FEC.Data[10100] := 286.55;
   Prof_FEC.Data[10101] := 318.04;
   Prof_FEC.Data[10102] := 341.41;
   Prof_FEC.Data[10103] := 358.64;
   Prof_FEC.Data[10104] := 409.95;
   Prof_FEC.Data[10105] := 421.98;
   Prof_FEC.Data[10106] := 432.22;
   Prof_FEC.Data[10107] := 458.88;
   Prof_FEC.Data[10108] := 467.71;
   Prof_FEC.Data[10109] := 535.09;
   Prof_FEC.Data[10110] := 509.99;
   Prof_FEC.Data[10111] := 555.36;
   Prof_FEC.Data[10112] := 560.54;
   Prof_FEC.Data[10113] := 591.59;
   Prof_FEC.Data[10114] := 634.12;
   Prof_FEC.Data[10115] := 664.87;
   Prof_FEC.Data[10116] := 596.51;
   Prof_FEC.Data[10117] := 657.79;
   Prof_FEC.Data[10118] := 655.76;
   Prof_FEC.Data[10119] := 615.66;
   Prof_FEC.Data[10120] := 591.8;
   Prof_FEC.Data[10121] := 691.74;
   Prof_FEC.Data[10122] := 622.02;
   Prof_FEC.Data[10123] := 692.4;
   Prof_FEC.Data[10124] := 625.57;
   Prof_FEC.Data[10125] := 645.69;
   Prof_FEC.Data[10126] := 625.76;
   Prof_FEC.Data[10127] := 608.64;
   Prof_FEC.Data[10128] := 576.09;
   Prof_FEC.Data[10129] := 580.63;
   Prof_FEC.Data[10130] := 726.57;
   Prof_FEC.Data[10131] := 560.89;
   Prof_FEC.Data[10132] := 559.26;
   Prof_FEC.Data[10133] := 643.29;
   Prof_FEC.Data[10134] := 575.18;
   Prof_FEC.Data[10135] := 602.17;
   Prof_FEC.Data[10136] := 575.39;
   Prof_FEC.Data[10137] := 689.5;
   Prof_FEC.Data[10138] := 617.81;
   Prof_FEC.Data[10139] := 707.53;
   Prof_FEC.Data[10140] := 732.67;
   Prof_FEC.Data[10141] := 775.66;
   Prof_FEC.Data[10142] := 723.22;
   Prof_FEC.Data[10143] := 582.77;
   Prof_FEC.Data[10144] := 304.25;
   Prof_FEC.Data[10145] := 180.62;
   Prof_FEC.Data[10146] := 119.85;
   Prof_FEC.Data[10147] := 116.35;
   Prof_FEC.Data[10148] := 86.39;
   Prof_FEC.Data[10149] := 56.62;
   Prof_FEC.Data[10150] := 58.26;
   Prof_FEC.Data[10151] := 59.91;
   Prof_FEC.Data[10152] := 92.46;
   Prof_FEC.Data[10153] := 97.38;
   Prof_FEC.Data[10154] := 127.49;
   Prof_FEC.Data[10155] := 139.0;
   Prof_FEC.Data[10156] := 33.172;
   Prof_FEC.Data[10157] := 35.364;
   Prof_FEC.Data[10158] := 34.306;
   Prof_FEC.Data[10159] := 36.232;
   Prof_FEC.Data[10160] := 34.174;
   Prof_FEC.Data[10161] := 34.383;
   Prof_FEC.Data[10162] := 33.423;
   Prof_FEC.Data[10163] := 34.235;
   Prof_FEC.Data[10164] := 35.554;
   Prof_FEC.Data[10165] := 32.183;
   Prof_FEC.Data[10166] := 33.496;
   Prof_FEC.Data[10167] := 33.543;
   Prof_FEC.Data[10168] := 34.615;
   Prof_FEC.Data[10169] := 36.921;
   Prof_FEC.Data[10170] := 37.924;
   Prof_FEC.Data[10171] := 35.111;
   Prof_FEC.Data[10172] := 37.399;
   Prof_FEC.Data[10173] := 35.343;
   Prof_FEC.Data[10174] := 35.173;
   Prof_FEC.Data[10175] := 36.576;
   Prof_FEC.Data[10176] := 37.03;
   Prof_FEC.Data[10177] := 35.161;
   Prof_FEC.Data[10178] := 36.066;
   Prof_FEC.Data[10179] := 35.318;
   Prof_FEC.Data[10180] := 36.244;
   Prof_FEC.Data[10181] := 35.315;
   Prof_FEC.Data[10182] := 36.693;
   Prof_FEC.Data[10183] := 33.878;
   Prof_FEC.Data[10184] := 35.225;
   Prof_FEC.Data[10185] := 34.875;
   Prof_FEC.Data[10186] := 34.406;
   Prof_FEC.Data[10187] := 32.983;
   Prof_FEC.Data[10188] := 34.195;
   Prof_FEC.Data[10189] := 33.546;
   Prof_FEC.Data[10190] := 33.016;
   Prof_FEC.Data[10191] := 34.941;
   Prof_FEC.Data[10192] := 32.475;
   Prof_FEC.Data[10193] := 32.511;
   Prof_FEC.Data[10194] := 32.755;
   Prof_FEC.Data[10195] := 35.676;
   Prof_FEC.Data[10196] := 236.9;
   Prof_FEC.Data[10197] := 282.32;
   Prof_FEC.Data[10198] := 273.33;
   Prof_FEC.Data[10199] := 330.07;
   Prof_FEC.Data[10200] := 373.3;
   Prof_FEC.Data[10201] := 348.52;
   Prof_FEC.Data[10202] := 367.36;
   Prof_FEC.Data[10203] := 378.71;
   Prof_FEC.Data[10204] := 470.3;
   Prof_FEC.Data[10205] := 447.66;
   Prof_FEC.Data[10206] := 497.43;
   Prof_FEC.Data[10207] := 504.23;
   Prof_FEC.Data[10208] := 592.0;
   Prof_FEC.Data[10209] := 648.79;
   Prof_FEC.Data[10210] := 581.1;
   Prof_FEC.Data[10211] := 599.12;
   Prof_FEC.Data[10212] := 599.89;
   Prof_FEC.Data[10213] := 537.75;
   Prof_FEC.Data[10214] := 609.71;
   Prof_FEC.Data[10215] := 586.59;
   Prof_FEC.Data[10216] := 621.68;
   Prof_FEC.Data[10217] := 589.59;
   Prof_FEC.Data[10218] := 569.5;
   Prof_FEC.Data[10219] := 530.8;
   Prof_FEC.Data[10220] := 573.79;
   Prof_FEC.Data[10221] := 502.16;
   Prof_FEC.Data[10222] := 610.83;
   Prof_FEC.Data[10223] := 550.59;
   Prof_FEC.Data[10224] := 545.7;
   Prof_FEC.Data[10225] := 532.09;
   Prof_FEC.Data[10226] := 599.05;
   Prof_FEC.Data[10227] := 571.08;
   Prof_FEC.Data[10228] := 590.8;
   Prof_FEC.Data[10229] := 661.3;
   Prof_FEC.Data[10230] := 639.43;
   Prof_FEC.Data[10231] := 627.3;
   Prof_FEC.Data[10232] := 637.87;
   Prof_FEC.Data[10233] := 627.85;
   Prof_FEC.Data[10234] := 571.66;
   Prof_FEC.Data[10235] := 652.21;
   Prof_FEC.Data[10236] := 659.57;
   Prof_FEC.Data[10237] := 732.98;
   Prof_FEC.Data[10238] := 645.06;
   Prof_FEC.Data[10239] := 528.42;
   Prof_FEC.Data[10240] := 250.36;
   Prof_FEC.Data[10241] := 157.88;
   Prof_FEC.Data[10242] := 119.5;
   Prof_FEC.Data[10243] := 103.41;
   Prof_FEC.Data[10244] := 75.98;
   Prof_FEC.Data[10245] := 54.98;
   Prof_FEC.Data[10246] := 45.22;
   Prof_FEC.Data[10247] := 61.57;
   Prof_FEC.Data[10248] := 85.88;
   Prof_FEC.Data[10249] := 107.39;
   Prof_FEC.Data[10250] := 114.12;
   Prof_FEC.Data[10251] := 135.66;
   Prof_FEC.Data[10252] := 33.375;
   Prof_FEC.Data[10253] := 33.688;
   Prof_FEC.Data[10254] := 34.315;
   Prof_FEC.Data[10255] := 35.025;
   Prof_FEC.Data[10256] := 34.414;
   Prof_FEC.Data[10257] := 36.052;
   Prof_FEC.Data[10258] := 34.805;
   Prof_FEC.Data[10259] := 34.895;
   Prof_FEC.Data[10260] := 34.573;
   Prof_FEC.Data[10261] := 31.169;
   Prof_FEC.Data[10262] := 30.591;
   Prof_FEC.Data[10263] := 32.24;
   Prof_FEC.Data[10264] := 37.132;
   Prof_FEC.Data[10265] := 35.119;
   Prof_FEC.Data[10266] := 34.158;
   Prof_FEC.Data[10267] := 35.458;
   Prof_FEC.Data[10268] := 32.155;
   Prof_FEC.Data[10269] := 32.767;
   Prof_FEC.Data[10270] := 34.818;
   Prof_FEC.Data[10271] := 33.785;
   Prof_FEC.Data[10272] := 34.577;
   Prof_FEC.Data[10273] := 35.015;
   Prof_FEC.Data[10274] := 35.168;
   Prof_FEC.Data[10275] := 34.406;
   Prof_FEC.Data[10276] := 34.486;
   Prof_FEC.Data[10277] := 35.279;
   Prof_FEC.Data[10278] := 33.354;
   Prof_FEC.Data[10279] := 35.397;
   Prof_FEC.Data[10280] := 36.398;
   Prof_FEC.Data[10281] := 37.425;
   Prof_FEC.Data[10282] := 37.721;
   Prof_FEC.Data[10283] := 36.888;
   Prof_FEC.Data[10284] := 33.938;
   Prof_FEC.Data[10285] := 34.307;
   Prof_FEC.Data[10286] := 36.249;
   Prof_FEC.Data[10287] := 35.981;
   Prof_FEC.Data[10288] := 35.442;
   Prof_FEC.Data[10289] := 35.023;
   Prof_FEC.Data[10290] := 38.749;
   Prof_FEC.Data[10291] := 39.029;
   Prof_FEC.Data[10292] := 289.41;
   Prof_FEC.Data[10293] := 313.54;
   Prof_FEC.Data[10294] := 329.73;
   Prof_FEC.Data[10295] := 321.57;
   Prof_FEC.Data[10296] := 368.03;
   Prof_FEC.Data[10297] := 390.9;
   Prof_FEC.Data[10298] := 480.31;
   Prof_FEC.Data[10299] := 466.2;
   Prof_FEC.Data[10300] := 469.87;
   Prof_FEC.Data[10301] := 565.88;
   Prof_FEC.Data[10302] := 526.33;
   Prof_FEC.Data[10303] := 611.2;
   Prof_FEC.Data[10304] := 676.9;
   Prof_FEC.Data[10305] := 726.17;
   Prof_FEC.Data[10306] := 698.13;
   Prof_FEC.Data[10307] := 737.54;
   Prof_FEC.Data[10308] := 691.91;
   Prof_FEC.Data[10309] := 758.7;
   Prof_FEC.Data[10310] := 700.33;
   Prof_FEC.Data[10311] := 773.9;
   Prof_FEC.Data[10312] := 764.79;
   Prof_FEC.Data[10313] := 745.05;
   Prof_FEC.Data[10314] := 680.56;
   Prof_FEC.Data[10315] := 716.2;
   Prof_FEC.Data[10316] := 658.72;
   Prof_FEC.Data[10317] := 539.44;
   Prof_FEC.Data[10318] := 612.1;
   Prof_FEC.Data[10319] := 653.96;
   Prof_FEC.Data[10320] := 684.64;
   Prof_FEC.Data[10321] := 723.99;
   Prof_FEC.Data[10322] := 749.77;
   Prof_FEC.Data[10323] := 684.87;
   Prof_FEC.Data[10324] := 602.76;
   Prof_FEC.Data[10325] := 658.51;
   Prof_FEC.Data[10326] := 664.29;
   Prof_FEC.Data[10327] := 609.6;
   Prof_FEC.Data[10328] := 621.7;
   Prof_FEC.Data[10329] := 599.78;
   Prof_FEC.Data[10330] := 605.82;
   Prof_FEC.Data[10331] := 561.66;
   Prof_FEC.Data[10332] := 685.09;
   Prof_FEC.Data[10333] := 673.12;
   Prof_FEC.Data[10334] := 599.78;
   Prof_FEC.Data[10335] := 509.49;
   Prof_FEC.Data[10336] := 275.34;
   Prof_FEC.Data[10337] := 197.32;
   Prof_FEC.Data[10338] := 120.34;
   Prof_FEC.Data[10339] := 108.34;
   Prof_FEC.Data[10340] := 79.39;
   Prof_FEC.Data[10341] := 63.99;
   Prof_FEC.Data[10342] := 59.08;
   Prof_FEC.Data[10343] := 67.65;
   Prof_FEC.Data[10344] := 96.89;
   Prof_FEC.Data[10345] := 101.61;
   Prof_FEC.Data[10346] := 128.04;
   Prof_FEC.Data[10347] := 141.98;
   Prof_FEC.Data[10348] := 33.78;
   Prof_FEC.Data[10349] := 35.267;
   Prof_FEC.Data[10350] := 36.15;
   Prof_FEC.Data[10351] := 35.848;
   Prof_FEC.Data[10352] := 35.786;
   Prof_FEC.Data[10353] := 36.559;
   Prof_FEC.Data[10354] := 36.169;
   Prof_FEC.Data[10355] := 38.093;
   Prof_FEC.Data[10356] := 37.72;
   Prof_FEC.Data[10357] := 35.855;
   Prof_FEC.Data[10358] := 35.224;
   Prof_FEC.Data[10359] := 34.212;
   Prof_FEC.Data[10360] := 35.207;
   Prof_FEC.Data[10361] := 34.734;
   Prof_FEC.Data[10362] := 35.007;
   Prof_FEC.Data[10363] := 35.016;
   Prof_FEC.Data[10364] := 32.835;
   Prof_FEC.Data[10365] := 31.919;
   Prof_FEC.Data[10366] := 33.853;
   Prof_FEC.Data[10367] := 33.766;
   Prof_FEC.Data[10368] := 34.723;
   Prof_FEC.Data[10369] := 34.23;
   Prof_FEC.Data[10370] := 35.056;
   Prof_FEC.Data[10371] := 35.157;
   Prof_FEC.Data[10372] := 35.14;
   Prof_FEC.Data[10373] := 35.786;
   Prof_FEC.Data[10374] := 35.289;
   Prof_FEC.Data[10375] := 37.409;
   Prof_FEC.Data[10376] := 37.081;
   Prof_FEC.Data[10377] := 36.531;
   Prof_FEC.Data[10378] := 35.831;
   Prof_FEC.Data[10379] := 38.461;
   Prof_FEC.Data[10380] := 37.536;
   Prof_FEC.Data[10381] := 35.133;
   Prof_FEC.Data[10382] := 36.709;
   Prof_FEC.Data[10383] := 36.354;
   Prof_FEC.Data[10384] := 38.088;
   Prof_FEC.Data[10385] := 38.974;
   Prof_FEC.Data[10386] := 36.905;
   Prof_FEC.Data[10387] := 34.615;
   Prof_FEC.Data[10388] := 127.6;
   Prof_FEC.Data[10389] := 115.12;
   Prof_FEC.Data[10390] := 114.94;
   Prof_FEC.Data[10391] := 151.84;
   Prof_FEC.Data[10392] := 212.95;
   Prof_FEC.Data[10393] := 276.19;
   Prof_FEC.Data[10394] := 318.55;
   Prof_FEC.Data[10395] := 312.22;
   Prof_FEC.Data[10396] := 277.77;
   Prof_FEC.Data[10397] := 294.54;
   Prof_FEC.Data[10398] := 316.43;
   Prof_FEC.Data[10399] := 294.57;
   Prof_FEC.Data[10400] := 349.95;
   Prof_FEC.Data[10401] := 386.2;
   Prof_FEC.Data[10402] := 357.1;
   Prof_FEC.Data[10403] := 393.85;
   Prof_FEC.Data[10404] := 387.49;
   Prof_FEC.Data[10405] := 375.2;
   Prof_FEC.Data[10406] := 375.23;
   Prof_FEC.Data[10407] := 318.82;
   Prof_FEC.Data[10408] := 350.91;
   Prof_FEC.Data[10409] := 366.82;
   Prof_FEC.Data[10410] := 342.53;
   Prof_FEC.Data[10411] := 326.85;
   Prof_FEC.Data[10412] := 229.79;
   Prof_FEC.Data[10413] := 267.44;
   Prof_FEC.Data[10414] := 250.87;
   Prof_FEC.Data[10415] := 251.8;
   Prof_FEC.Data[10416] := 299.96;
   Prof_FEC.Data[10417] := 287.53;
   Prof_FEC.Data[10418] := 261.77;
   Prof_FEC.Data[10419] := 275.38;
   Prof_FEC.Data[10420] := 265.69;
   Prof_FEC.Data[10421] := 253.09;
   Prof_FEC.Data[10422] := 280.67;
   Prof_FEC.Data[10423] := 254.2;
   Prof_FEC.Data[10424] := 308.94;
   Prof_FEC.Data[10425] := 313.94;
   Prof_FEC.Data[10426] := 299.08;
   Prof_FEC.Data[10427] := 228.47;
   Prof_FEC.Data[10428] := 89.78;
   Prof_FEC.Data[10429] := 54.77;
   Prof_FEC.Data[10430] := 36.33;
   Prof_FEC.Data[10431] := 35.62;
   Prof_FEC.Data[10432] := 51.17;
   Prof_FEC.Data[10433] := 56.05;
   Prof_FEC.Data[10434] := 50.38;
   Prof_FEC.Data[10435] := 52.86;
   Prof_FEC.Data[10436] := 46.89;
   Prof_FEC.Data[10437] := 49.85;
   Prof_FEC.Data[10438] := 51.46;
   Prof_FEC.Data[10439] := 53.88;
   Prof_FEC.Data[10440] := 54.56;
   Prof_FEC.Data[10441] := 60.36;
   Prof_FEC.Data[10442] := 70.92;
   Prof_FEC.Data[10443] := 90.73;
   Prof_FEC.Data[10444] := 31.108;
   Prof_FEC.Data[10445] := 34.284;
   Prof_FEC.Data[10446] := 33.876;
   Prof_FEC.Data[10447] := 31.209;
   Prof_FEC.Data[10448] := 31.951;
   Prof_FEC.Data[10449] := 32.206;
   Prof_FEC.Data[10450] := 30.333;
   Prof_FEC.Data[10451] := 30.849;
   Prof_FEC.Data[10452] := 33.682;
   Prof_FEC.Data[10453] := 34.985;
   Prof_FEC.Data[10454] := 35.462;
   Prof_FEC.Data[10455] := 34.687;
   Prof_FEC.Data[10456] := 35.945;
   Prof_FEC.Data[10457] := 32.596;
   Prof_FEC.Data[10458] := 32.374;
   Prof_FEC.Data[10459] := 31.772;
   Prof_FEC.Data[10460] := 32.471;
   Prof_FEC.Data[10461] := 34.415;
   Prof_FEC.Data[10462] := 36.665;
   Prof_FEC.Data[10463] := 34.693;
   Prof_FEC.Data[10464] := 34.714;
   Prof_FEC.Data[10465] := 34.342;
   Prof_FEC.Data[10466] := 34.757;
   Prof_FEC.Data[10467] := 33.885;
   Prof_FEC.Data[10468] := 35.648;
   Prof_FEC.Data[10469] := 32.64;
   Prof_FEC.Data[10470] := 35.206;
   Prof_FEC.Data[10471] := 35.741;
   Prof_FEC.Data[10472] := 34.625;
   Prof_FEC.Data[10473] := 33.011;
   Prof_FEC.Data[10474] := 31.987;
   Prof_FEC.Data[10475] := 32.246;
   Prof_FEC.Data[10476] := 33.409;
   Prof_FEC.Data[10477] := 34.593;
   Prof_FEC.Data[10478] := 35.015;
   Prof_FEC.Data[10479] := 34.623;
   Prof_FEC.Data[10480] := 36.369;
   Prof_FEC.Data[10481] := 35.349;
   Prof_FEC.Data[10482] := 35.031;
   Prof_FEC.Data[10483] := 33.136;
   Prof_FEC.Data[10484] := 158.18;
   Prof_FEC.Data[10485] := 122.93;
   Prof_FEC.Data[10486] := 115.22;
   Prof_FEC.Data[10487] := 99.26;
   Prof_FEC.Data[10488] := 79.21;
   Prof_FEC.Data[10489] := 62.24;
   Prof_FEC.Data[10490] := 61.16;
   Prof_FEC.Data[10491] := 57.6;
   Prof_FEC.Data[10492] := 76.41;
   Prof_FEC.Data[10493] := 79.74;
   Prof_FEC.Data[10494] := 81.15;
   Prof_FEC.Data[10495] := 73.02;
   Prof_FEC.Data[10496] := 75.9;
   Prof_FEC.Data[10497] := 68.97;
   Prof_FEC.Data[10498] := 62.9;
   Prof_FEC.Data[10499] := 69.8;
   Prof_FEC.Data[10500] := 74.07;
   Prof_FEC.Data[10501] := 75.53;
   Prof_FEC.Data[10502] := 75.7;
   Prof_FEC.Data[10503] := 72.23;
   Prof_FEC.Data[10504] := 63.42;
   Prof_FEC.Data[10505] := 72.83;
   Prof_FEC.Data[10506] := 60.55;
   Prof_FEC.Data[10507] := 66.45;
   Prof_FEC.Data[10508] := 68.43;
   Prof_FEC.Data[10509] := 64.92;
   Prof_FEC.Data[10510] := 63.28;
   Prof_FEC.Data[10511] := 63.68;
   Prof_FEC.Data[10512] := 64.25;
   Prof_FEC.Data[10513] := 60.53;
   Prof_FEC.Data[10514] := 63.28;
   Prof_FEC.Data[10515] := 58.41;
   Prof_FEC.Data[10516] := 65.86;
   Prof_FEC.Data[10517] := 66.56;
   Prof_FEC.Data[10518] := 70.14;
   Prof_FEC.Data[10519] := 66.02;
   Prof_FEC.Data[10520] := 62.91;
   Prof_FEC.Data[10521] := 60.76;
   Prof_FEC.Data[10522] := 61.19;
   Prof_FEC.Data[10523] := 59.9;
   Prof_FEC.Data[10524] := 70.71;
   Prof_FEC.Data[10525] := 75.38;
   Prof_FEC.Data[10526] := 83.37;
   Prof_FEC.Data[10527] := 71.69;
   Prof_FEC.Data[10528] := 70.9;
   Prof_FEC.Data[10529] := 65.59;
   Prof_FEC.Data[10530] := 64.11;
   Prof_FEC.Data[10531] := 78.17;
   Prof_FEC.Data[10532] := 87.17;
   Prof_FEC.Data[10533] := 84.83;
   Prof_FEC.Data[10534] := 82.21;
   Prof_FEC.Data[10535] := 93.06;
   Prof_FEC.Data[10536] := 86.63;
   Prof_FEC.Data[10537] := 99.34;
   Prof_FEC.Data[10538] := 109.36;
   Prof_FEC.Data[10539] := 130.9;
   Prof_FEC.Data[10540] := 37.245;
   Prof_FEC.Data[10541] := 40.299;
   Prof_FEC.Data[10542] := 41.773;
   Prof_FEC.Data[10543] := 41.354;
   Prof_FEC.Data[10544] := 38.723;
   Prof_FEC.Data[10545] := 37.341;
   Prof_FEC.Data[10546] := 36.573;
   Prof_FEC.Data[10547] := 36.094;
   Prof_FEC.Data[10548] := 37.229;
   Prof_FEC.Data[10549] := 37.337;
   Prof_FEC.Data[10550] := 36.757;
   Prof_FEC.Data[10551] := 35.936;
   Prof_FEC.Data[10552] := 35.259;
   Prof_FEC.Data[10553] := 34.958;
   Prof_FEC.Data[10554] := 33.232;
   Prof_FEC.Data[10555] := 36.206;
   Prof_FEC.Data[10556] := 36.113;
   Prof_FEC.Data[10557] := 34.954;
   Prof_FEC.Data[10558] := 36.995;
   Prof_FEC.Data[10559] := 34.302;
   Prof_FEC.Data[10560] := 33.61;
   Prof_FEC.Data[10561] := 34.085;
   Prof_FEC.Data[10562] := 35.509;
   Prof_FEC.Data[10563] := 33.865;
   Prof_FEC.Data[10564] := 33.368;
   Prof_FEC.Data[10565] := 34.167;
   Prof_FEC.Data[10566] := 36.295;
   Prof_FEC.Data[10567] := 35.915;
   Prof_FEC.Data[10568] := 35.04;
   Prof_FEC.Data[10569] := 34.085;
   Prof_FEC.Data[10570] := 35.162;
   Prof_FEC.Data[10571] := 36.035;
   Prof_FEC.Data[10572] := 33.567;
   Prof_FEC.Data[10573] := 37.904;
   Prof_FEC.Data[10574] := 36.252;
   Prof_FEC.Data[10575] := 39.589;
   Prof_FEC.Data[10576] := 33.685;
   Prof_FEC.Data[10577] := 34.946;
   Prof_FEC.Data[10578] := 35.395;
   Prof_FEC.Data[10579] := 39.064;
   Prof_FEC.Data[10580] := 286.01;
   Prof_FEC.Data[10581] := 307.42;
   Prof_FEC.Data[10582] := 342.11;
   Prof_FEC.Data[10583] := 345.28;
   Prof_FEC.Data[10584] := 348.38;
   Prof_FEC.Data[10585] := 408.54;
   Prof_FEC.Data[10586] := 411.6;
   Prof_FEC.Data[10587] := 419.11;
   Prof_FEC.Data[10588] := 458.83;
   Prof_FEC.Data[10589] := 519.87;
   Prof_FEC.Data[10590] := 516.19;
   Prof_FEC.Data[10591] := 596.15;
   Prof_FEC.Data[10592] := 583.47;
   Prof_FEC.Data[10593] := 635.02;
   Prof_FEC.Data[10594] := 651.21;
   Prof_FEC.Data[10595] := 571.17;
   Prof_FEC.Data[10596] := 553.11;
   Prof_FEC.Data[10597] := 621.24;
   Prof_FEC.Data[10598] := 635.9;
   Prof_FEC.Data[10599] := 613.61;
   Prof_FEC.Data[10600] := 594.43;
   Prof_FEC.Data[10601] := 554.95;
   Prof_FEC.Data[10602] := 575.17;
   Prof_FEC.Data[10603] := 581.45;
   Prof_FEC.Data[10604] := 545.71;
   Prof_FEC.Data[10605] := 558.33;
   Prof_FEC.Data[10606] := 607.89;
   Prof_FEC.Data[10607] := 589.02;
   Prof_FEC.Data[10608] := 645.38;
   Prof_FEC.Data[10609] := 661.8;
   Prof_FEC.Data[10610] := 626.51;
   Prof_FEC.Data[10611] := 602.56;
   Prof_FEC.Data[10612] := 608.16;
   Prof_FEC.Data[10613] := 612.47;
   Prof_FEC.Data[10614] := 652.81;
   Prof_FEC.Data[10615] := 624.17;
   Prof_FEC.Data[10616] := 647.64;
   Prof_FEC.Data[10617] := 655.72;
   Prof_FEC.Data[10618] := 666.43;
   Prof_FEC.Data[10619] := 627.8;
   Prof_FEC.Data[10620] := 715.02;
   Prof_FEC.Data[10621] := 738.41;
   Prof_FEC.Data[10622] := 671.43;
   Prof_FEC.Data[10623] := 582.69;
   Prof_FEC.Data[10624] := 286.65;
   Prof_FEC.Data[10625] := 209.91;
   Prof_FEC.Data[10626] := 139.29;
   Prof_FEC.Data[10627] := 118.15;
   Prof_FEC.Data[10628] := 102.76;
   Prof_FEC.Data[10629] := 79.2;
   Prof_FEC.Data[10630] := 62.53;
   Prof_FEC.Data[10631] := 78.59;
   Prof_FEC.Data[10632] := 94.33;
   Prof_FEC.Data[10633] := 99.84;
   Prof_FEC.Data[10634] := 118.34;
   Prof_FEC.Data[10635] := 127.79;
   Prof_FEC.Data[10636] := 33.982;
   Prof_FEC.Data[10637] := 35.7;
   Prof_FEC.Data[10638] := 40.87;
   Prof_FEC.Data[10639] := 40.205;
   Prof_FEC.Data[10640] := 39.055;
   Prof_FEC.Data[10641] := 39.436;
   Prof_FEC.Data[10642] := 40.58;
   Prof_FEC.Data[10643] := 39.541;
   Prof_FEC.Data[10644] := 37.886;
   Prof_FEC.Data[10645] := 38.012;
   Prof_FEC.Data[10646] := 37.734;
   Prof_FEC.Data[10647] := 37.225;
   Prof_FEC.Data[10648] := 38.033;
   Prof_FEC.Data[10649] := 38.761;
   Prof_FEC.Data[10650] := 38.047;
   Prof_FEC.Data[10651] := 37.506;
   Prof_FEC.Data[10652] := 39.05;
   Prof_FEC.Data[10653] := 37.604;
   Prof_FEC.Data[10654] := 38.674;
   Prof_FEC.Data[10655] := 36.61;
   Prof_FEC.Data[10656] := 40.26;
   Prof_FEC.Data[10657] := 38.905;
   Prof_FEC.Data[10658] := 39.885;
   Prof_FEC.Data[10659] := 39.231;
   Prof_FEC.Data[10660] := 39.343;
   Prof_FEC.Data[10661] := 38.045;
   Prof_FEC.Data[10662] := 35.682;
   Prof_FEC.Data[10663] := 38.328;
   Prof_FEC.Data[10664] := 38.153;
   Prof_FEC.Data[10665] := 38.891;
   Prof_FEC.Data[10666] := 38.659;
   Prof_FEC.Data[10667] := 38.714;
   Prof_FEC.Data[10668] := 37.522;
   Prof_FEC.Data[10669] := 35.329;
   Prof_FEC.Data[10670] := 37.55;
   Prof_FEC.Data[10671] := 38.702;
   Prof_FEC.Data[10672] := 38.811;
   Prof_FEC.Data[10673] := 40.505;
   Prof_FEC.Data[10674] := 41.996;
   Prof_FEC.Data[10675] := 43.019;
   Prof_FEC.Data[10676] := 349.57;
   Prof_FEC.Data[10677] := 326.08;
   Prof_FEC.Data[10678] := 351.61;
   Prof_FEC.Data[10679] := 368.81;
   Prof_FEC.Data[10680] := 379.27;
   Prof_FEC.Data[10681] := 395.95;
   Prof_FEC.Data[10682] := 461.22;
   Prof_FEC.Data[10683] := 486.95;
   Prof_FEC.Data[10684] := 502.31;
   Prof_FEC.Data[10685] := 584.58;
   Prof_FEC.Data[10686] := 607.45;
   Prof_FEC.Data[10687] := 532.19;
   Prof_FEC.Data[10688] := 665.69;
   Prof_FEC.Data[10689] := 682.17;
   Prof_FEC.Data[10690] := 674.4;
   Prof_FEC.Data[10691] := 679.38;
   Prof_FEC.Data[10692] := 536.5;
   Prof_FEC.Data[10693] := 609.12;
   Prof_FEC.Data[10694] := 656.33;
   Prof_FEC.Data[10695] := 604.67;
   Prof_FEC.Data[10696] := 632.88;
   Prof_FEC.Data[10697] := 682.73;
   Prof_FEC.Data[10698] := 633.51;
   Prof_FEC.Data[10699] := 577.52;
   Prof_FEC.Data[10700] := 603.91;
   Prof_FEC.Data[10701] := 528.61;
   Prof_FEC.Data[10702] := 606.85;
   Prof_FEC.Data[10703] := 634.34;
   Prof_FEC.Data[10704] := 644.82;
   Prof_FEC.Data[10705] := 682.18;
   Prof_FEC.Data[10706] := 676.87;
   Prof_FEC.Data[10707] := 695.3;
   Prof_FEC.Data[10708] := 762.79;
   Prof_FEC.Data[10709] := 643.86;
   Prof_FEC.Data[10710] := 744.4;
   Prof_FEC.Data[10711] := 730.47;
   Prof_FEC.Data[10712] := 696.8;
   Prof_FEC.Data[10713] := 651.16;
   Prof_FEC.Data[10714] := 690.98;
   Prof_FEC.Data[10715] := 662.25;
   Prof_FEC.Data[10716] := 727.58;
   Prof_FEC.Data[10717] := 768.22;
   Prof_FEC.Data[10718] := 664.91;
   Prof_FEC.Data[10719] := 537.17;
   Prof_FEC.Data[10720] := 272.76;
   Prof_FEC.Data[10721] := 201.22;
   Prof_FEC.Data[10722] := 146.25;
   Prof_FEC.Data[10723] := 121.39;
   Prof_FEC.Data[10724] := 88.32;
   Prof_FEC.Data[10725] := 67.61;
   Prof_FEC.Data[10726] := 66.78;
   Prof_FEC.Data[10727] := 73.9;
   Prof_FEC.Data[10728] := 89.09;
   Prof_FEC.Data[10729] := 100.83;
   Prof_FEC.Data[10730] := 110.82;
   Prof_FEC.Data[10731] := 115.51;
   Prof_FEC.Data[10732] := 33.347;
   Prof_FEC.Data[10733] := 34.606;
   Prof_FEC.Data[10734] := 36.162;
   Prof_FEC.Data[10735] := 35.586;
   Prof_FEC.Data[10736] := 35.616;
   Prof_FEC.Data[10737] := 35.052;
   Prof_FEC.Data[10738] := 34.457;
   Prof_FEC.Data[10739] := 37.098;
   Prof_FEC.Data[10740] := 31.835;
   Prof_FEC.Data[10741] := 33.109;
   Prof_FEC.Data[10742] := 34.521;
   Prof_FEC.Data[10743] := 35.657;
   Prof_FEC.Data[10744] := 34.363;
   Prof_FEC.Data[10745] := 34.324;
   Prof_FEC.Data[10746] := 35.778;
   Prof_FEC.Data[10747] := 36.336;
   Prof_FEC.Data[10748] := 33.605;
   Prof_FEC.Data[10749] := 33.398;
   Prof_FEC.Data[10750] := 35.04;
   Prof_FEC.Data[10751] := 37.15;
   Prof_FEC.Data[10752] := 36.831;
   Prof_FEC.Data[10753] := 38.128;
   Prof_FEC.Data[10754] := 39.053;
   Prof_FEC.Data[10755] := 39.527;
   Prof_FEC.Data[10756] := 35.998;
   Prof_FEC.Data[10757] := 36.653;
   Prof_FEC.Data[10758] := 39.425;
   Prof_FEC.Data[10759] := 37.127;
   Prof_FEC.Data[10760] := 38.596;
   Prof_FEC.Data[10761] := 39.711;
   Prof_FEC.Data[10762] := 41.74;
   Prof_FEC.Data[10763] := 39.526;
   Prof_FEC.Data[10764] := 38.12;
   Prof_FEC.Data[10765] := 34.444;
   Prof_FEC.Data[10766] := 38.218;
   Prof_FEC.Data[10767] := 36.412;
   Prof_FEC.Data[10768] := 40.861;
   Prof_FEC.Data[10769] := 40.611;
   Prof_FEC.Data[10770] := 38.708;
   Prof_FEC.Data[10771] := 37.987;
   Prof_FEC.Data[10772] := 278.27;
   Prof_FEC.Data[10773] := 325.22;
   Prof_FEC.Data[10774] := 347.56;
   Prof_FEC.Data[10775] := 399.25;
   Prof_FEC.Data[10776] := 397.72;
   Prof_FEC.Data[10777] := 464.36;
   Prof_FEC.Data[10778] := 414.47;
   Prof_FEC.Data[10779] := 466.49;
   Prof_FEC.Data[10780] := 499.69;
   Prof_FEC.Data[10781] := 593.51;
   Prof_FEC.Data[10782] := 565.77;
   Prof_FEC.Data[10783] := 666.65;
   Prof_FEC.Data[10784] := 650.18;
   Prof_FEC.Data[10785] := 634.17;
   Prof_FEC.Data[10786] := 631.15;
   Prof_FEC.Data[10787] := 572.64;
   Prof_FEC.Data[10788] := 613.22;
   Prof_FEC.Data[10789] := 574.28;
   Prof_FEC.Data[10790] := 647.05;
   Prof_FEC.Data[10791] := 675.94;
   Prof_FEC.Data[10792] := 646.02;
   Prof_FEC.Data[10793] := 705.6;
   Prof_FEC.Data[10794] := 651.31;
   Prof_FEC.Data[10795] := 655.54;
   Prof_FEC.Data[10796] := 581.23;
   Prof_FEC.Data[10797] := 610.54;
   Prof_FEC.Data[10798] := 605.16;
   Prof_FEC.Data[10799] := 645.29;
   Prof_FEC.Data[10800] := 588.65;
   Prof_FEC.Data[10801] := 627.93;
   Prof_FEC.Data[10802] := 566.23;
   Prof_FEC.Data[10803] := 600.94;
   Prof_FEC.Data[10804] := 575.05;
   Prof_FEC.Data[10805] := 550.26;
   Prof_FEC.Data[10806] := 581.76;
   Prof_FEC.Data[10807] := 609.23;
   Prof_FEC.Data[10808] := 569.87;
   Prof_FEC.Data[10809] := 586.61;
   Prof_FEC.Data[10810] := 635.55;
   Prof_FEC.Data[10811] := 628.98;
   Prof_FEC.Data[10812] := 658.75;
   Prof_FEC.Data[10813] := 691.3;
   Prof_FEC.Data[10814] := 669.93;
   Prof_FEC.Data[10815] := 524.5;
   Prof_FEC.Data[10816] := 294.78;
   Prof_FEC.Data[10817] := 187.24;
   Prof_FEC.Data[10818] := 120.34;
   Prof_FEC.Data[10819] := 94.93;
   Prof_FEC.Data[10820] := 80.03;
   Prof_FEC.Data[10821] := 51.21;
   Prof_FEC.Data[10822] := 51.54;
   Prof_FEC.Data[10823] := 49.53;
   Prof_FEC.Data[10824] := 74.95;
   Prof_FEC.Data[10825] := 81.75;
   Prof_FEC.Data[10826] := 102.03;
   Prof_FEC.Data[10827] := 112.51;
   Prof_FEC.Data[10828] := 30.465;
   Prof_FEC.Data[10829] := 33.692;
   Prof_FEC.Data[10830] := 33.765;
   Prof_FEC.Data[10831] := 35.875;
   Prof_FEC.Data[10832] := 35.675;
   Prof_FEC.Data[10833] := 35.506;
   Prof_FEC.Data[10834] := 35.127;
   Prof_FEC.Data[10835] := 35.153;
   Prof_FEC.Data[10836] := 35.024;
   Prof_FEC.Data[10837] := 33.814;
   Prof_FEC.Data[10838] := 34.43;
   Prof_FEC.Data[10839] := 34.351;
   Prof_FEC.Data[10840] := 36.262;
   Prof_FEC.Data[10841] := 36.805;
   Prof_FEC.Data[10842] := 38.3;
   Prof_FEC.Data[10843] := 38.414;
   Prof_FEC.Data[10844] := 38.133;
   Prof_FEC.Data[10845] := 37.285;
   Prof_FEC.Data[10846] := 37.445;
   Prof_FEC.Data[10847] := 38.83;
   Prof_FEC.Data[10848] := 37.756;
   Prof_FEC.Data[10849] := 40.571;
   Prof_FEC.Data[10850] := 40.541;
   Prof_FEC.Data[10851] := 40.835;
   Prof_FEC.Data[10852] := 38.71;
   Prof_FEC.Data[10853] := 39.164;
   Prof_FEC.Data[10854] := 39.292;
   Prof_FEC.Data[10855] := 37.572;
   Prof_FEC.Data[10856] := 40.645;
   Prof_FEC.Data[10857] := 39.278;
   Prof_FEC.Data[10858] := 40.564;
   Prof_FEC.Data[10859] := 38.817;
   Prof_FEC.Data[10860] := 36.579;
   Prof_FEC.Data[10861] := 36.342;
   Prof_FEC.Data[10862] := 37.443;
   Prof_FEC.Data[10863] := 37.143;
   Prof_FEC.Data[10864] := 36.632;
   Prof_FEC.Data[10865] := 38.614;
   Prof_FEC.Data[10866] := 40.319;
   Prof_FEC.Data[10867] := 40.934;
   Prof_FEC.Data[10868] := 246.83;
   Prof_FEC.Data[10869] := 296.89;
   Prof_FEC.Data[10870] := 335.56;
   Prof_FEC.Data[10871] := 367.3;
   Prof_FEC.Data[10872] := 432.83;
   Prof_FEC.Data[10873] := 445.4;
   Prof_FEC.Data[10874] := 485.45;
   Prof_FEC.Data[10875] := 513.59;
   Prof_FEC.Data[10876] := 569.62;
   Prof_FEC.Data[10877] := 604.26;
   Prof_FEC.Data[10878] := 607.31;
   Prof_FEC.Data[10879] := 655.87;
   Prof_FEC.Data[10880] := 603.47;
   Prof_FEC.Data[10881] := 659.07;
   Prof_FEC.Data[10882] := 673.04;
   Prof_FEC.Data[10883] := 637.77;
   Prof_FEC.Data[10884] := 628.95;
   Prof_FEC.Data[10885] := 644.81;
   Prof_FEC.Data[10886] := 671.7;
   Prof_FEC.Data[10887] := 643.16;
   Prof_FEC.Data[10888] := 646.37;
   Prof_FEC.Data[10889] := 673.74;
   Prof_FEC.Data[10890] := 608.4;
   Prof_FEC.Data[10891] := 700.62;
   Prof_FEC.Data[10892] := 603.42;
   Prof_FEC.Data[10893] := 648.04;
   Prof_FEC.Data[10894] := 650.68;
   Prof_FEC.Data[10895] := 683.88;
   Prof_FEC.Data[10896] := 714.96;
   Prof_FEC.Data[10897] := 696.54;
   Prof_FEC.Data[10898] := 715.97;
   Prof_FEC.Data[10899] := 691.59;
   Prof_FEC.Data[10900] := 623.94;
   Prof_FEC.Data[10901] := 628.48;
   Prof_FEC.Data[10902] := 603.85;
   Prof_FEC.Data[10903] := 613.61;
   Prof_FEC.Data[10904] := 649.87;
   Prof_FEC.Data[10905] := 707.15;
   Prof_FEC.Data[10906] := 591.35;
   Prof_FEC.Data[10907] := 642.98;
   Prof_FEC.Data[10908] := 776.49;
   Prof_FEC.Data[10909] := 751.57;
   Prof_FEC.Data[10910] := 671.11;
   Prof_FEC.Data[10911] := 460.81;
   Prof_FEC.Data[10912] := 284.42;
   Prof_FEC.Data[10913] := 187.27;
   Prof_FEC.Data[10914] := 129.96;
   Prof_FEC.Data[10915] := 102.87;
   Prof_FEC.Data[10916] := 93.84;
   Prof_FEC.Data[10917] := 61.51;
   Prof_FEC.Data[10918] := 54.44;
   Prof_FEC.Data[10919] := 69.36;
   Prof_FEC.Data[10920] := 85.57;
   Prof_FEC.Data[10921] := 84.05;
   Prof_FEC.Data[10922] := 94.05;
   Prof_FEC.Data[10923] := 113.08;
   Prof_FEC.Data[10924] := 31.865;
   Prof_FEC.Data[10925] := 32.219;
   Prof_FEC.Data[10926] := 35.801;
   Prof_FEC.Data[10927] := 34.662;
   Prof_FEC.Data[10928] := 34.678;
   Prof_FEC.Data[10929] := 33.236;
   Prof_FEC.Data[10930] := 35.262;
   Prof_FEC.Data[10931] := 35.665;
   Prof_FEC.Data[10932] := 32.377;
   Prof_FEC.Data[10933] := 32.465;
   Prof_FEC.Data[10934] := 32.497;
   Prof_FEC.Data[10935] := 32.743;
   Prof_FEC.Data[10936] := 34.744;
   Prof_FEC.Data[10937] := 34.037;
   Prof_FEC.Data[10938] := 35.132;
   Prof_FEC.Data[10939] := 34.259;
   Prof_FEC.Data[10940] := 33.88;
   Prof_FEC.Data[10941] := 34.242;
   Prof_FEC.Data[10942] := 32.315;
   Prof_FEC.Data[10943] := 32.981;
   Prof_FEC.Data[10944] := 32.531;
   Prof_FEC.Data[10945] := 34.061;
   Prof_FEC.Data[10946] := 33.381;
   Prof_FEC.Data[10947] := 34.355;
   Prof_FEC.Data[10948] := 32.585;
   Prof_FEC.Data[10949] := 32.423;
   Prof_FEC.Data[10950] := 32.556;
   Prof_FEC.Data[10951] := 34.272;
   Prof_FEC.Data[10952] := 32.38;
   Prof_FEC.Data[10953] := 34.775;
   Prof_FEC.Data[10954] := 33.585;
   Prof_FEC.Data[10955] := 31.852;
   Prof_FEC.Data[10956] := 35.789;
   Prof_FEC.Data[10957] := 33.119;
   Prof_FEC.Data[10958] := 32.849;
   Prof_FEC.Data[10959] := 31.61;
   Prof_FEC.Data[10960] := 33.49;
   Prof_FEC.Data[10961] := 34.742;
   Prof_FEC.Data[10962] := 35.855;
   Prof_FEC.Data[10963] := 36.386;
   Prof_FEC.Data[10964] := 249.74;
   Prof_FEC.Data[10965] := 288.85;
   Prof_FEC.Data[10966] := 309.05;
   Prof_FEC.Data[10967] := 356.08;
   Prof_FEC.Data[10968] := 422.19;
   Prof_FEC.Data[10969] := 447.18;
   Prof_FEC.Data[10970] := 502.26;
   Prof_FEC.Data[10971] := 484.15;
   Prof_FEC.Data[10972] := 546.99;
   Prof_FEC.Data[10973] := 585.72;
   Prof_FEC.Data[10974] := 513.2;
   Prof_FEC.Data[10975] := 605.66;
   Prof_FEC.Data[10976] := 620.96;
   Prof_FEC.Data[10977] := 640.33;
   Prof_FEC.Data[10978] := 653.95;
   Prof_FEC.Data[10979] := 656.11;
   Prof_FEC.Data[10980] := 596.43;
   Prof_FEC.Data[10981] := 644.99;
   Prof_FEC.Data[10982] := 646.39;
   Prof_FEC.Data[10983] := 698.89;
   Prof_FEC.Data[10984] := 671.61;
   Prof_FEC.Data[10985] := 704.97;
   Prof_FEC.Data[10986] := 676.13;
   Prof_FEC.Data[10987] := 641.96;
   Prof_FEC.Data[10988] := 649.7;
   Prof_FEC.Data[10989] := 672.55;
   Prof_FEC.Data[10990] := 625.62;
   Prof_FEC.Data[10991] := 645.27;
   Prof_FEC.Data[10992] := 717.01;
   Prof_FEC.Data[10993] := 662.62;
   Prof_FEC.Data[10994] := 662.58;
   Prof_FEC.Data[10995] := 708.23;
   Prof_FEC.Data[10996] := 704.32;
   Prof_FEC.Data[10997] := 648.43;
   Prof_FEC.Data[10998] := 785.88;
   Prof_FEC.Data[10999] := 650.39;
   Prof_FEC.Data[11000] := 686.21;
   Prof_FEC.Data[11001] := 620.12;
   Prof_FEC.Data[11002] := 735.27;
   Prof_FEC.Data[11003] := 663.89;
   Prof_FEC.Data[11004] := 723.45;
   Prof_FEC.Data[11005] := 664.64;
   Prof_FEC.Data[11006] := 751.04;
   Prof_FEC.Data[11007] := 543.21;
   Prof_FEC.Data[11008] := 293.14;
   Prof_FEC.Data[11009] := 199.48;
   Prof_FEC.Data[11010] := 137.69;
   Prof_FEC.Data[11011] := 105.39;
   Prof_FEC.Data[11012] := 92.12;
   Prof_FEC.Data[11013] := 72.55;
   Prof_FEC.Data[11014] := 67.68;
   Prof_FEC.Data[11015] := 78.16;
   Prof_FEC.Data[11016] := 92.51;
   Prof_FEC.Data[11017] := 111.46;
   Prof_FEC.Data[11018] := 121.63;
   Prof_FEC.Data[11019] := 134.87;
   Prof_FEC.Data[11020] := 33.486;
   Prof_FEC.Data[11021] := 36.535;
   Prof_FEC.Data[11022] := 39.129;
   Prof_FEC.Data[11023] := 39.846;
   Prof_FEC.Data[11024] := 38.135;
   Prof_FEC.Data[11025] := 42.255;
   Prof_FEC.Data[11026] := 39.994;
   Prof_FEC.Data[11027] := 39.415;
   Prof_FEC.Data[11028] := 37.663;
   Prof_FEC.Data[11029] := 38.709;
   Prof_FEC.Data[11030] := 38.361;
   Prof_FEC.Data[11031] := 37.806;
   Prof_FEC.Data[11032] := 40.207;
   Prof_FEC.Data[11033] := 38.622;
   Prof_FEC.Data[11034] := 38.338;
   Prof_FEC.Data[11035] := 37.469;
   Prof_FEC.Data[11036] := 36.764;
   Prof_FEC.Data[11037] := 36.32;
   Prof_FEC.Data[11038] := 37.28;
   Prof_FEC.Data[11039] := 37.358;
   Prof_FEC.Data[11040] := 40.812;
   Prof_FEC.Data[11041] := 40.224;
   Prof_FEC.Data[11042] := 41.801;
   Prof_FEC.Data[11043] := 39.974;
   Prof_FEC.Data[11044] := 39.79;
   Prof_FEC.Data[11045] := 39.399;
   Prof_FEC.Data[11046] := 39.618;
   Prof_FEC.Data[11047] := 38.885;
   Prof_FEC.Data[11048] := 38.226;
   Prof_FEC.Data[11049] := 40.132;
   Prof_FEC.Data[11050] := 37.869;
   Prof_FEC.Data[11051] := 37.7;
   Prof_FEC.Data[11052] := 38.954;
   Prof_FEC.Data[11053] := 40.299;
   Prof_FEC.Data[11054] := 38.314;
   Prof_FEC.Data[11055] := 39.756;
   Prof_FEC.Data[11056] := 40.712;
   Prof_FEC.Data[11057] := 41.921;
   Prof_FEC.Data[11058] := 38.98;
   Prof_FEC.Data[11059] := 35.298;
   Prof_FEC.Data[11060] := 128.3;
   Prof_FEC.Data[11061] := 111.13;
   Prof_FEC.Data[11062] := 111.67;
   Prof_FEC.Data[11063] := 136.53;
   Prof_FEC.Data[11064] := 208.57;
   Prof_FEC.Data[11065] := 302.32;
   Prof_FEC.Data[11066] := 327.93;
   Prof_FEC.Data[11067] := 292.06;
   Prof_FEC.Data[11068] := 292.78;
   Prof_FEC.Data[11069] := 294.53;
   Prof_FEC.Data[11070] := 313.84;
   Prof_FEC.Data[11071] := 305.7;
   Prof_FEC.Data[11072] := 340.04;
   Prof_FEC.Data[11073] := 334.92;
   Prof_FEC.Data[11074] := 355.08;
   Prof_FEC.Data[11075] := 375.71;
   Prof_FEC.Data[11076] := 381.4;
   Prof_FEC.Data[11077] := 356.19;
   Prof_FEC.Data[11078] := 398.86;
   Prof_FEC.Data[11079] := 370.56;
   Prof_FEC.Data[11080] := 360.31;
   Prof_FEC.Data[11081] := 403.56;
   Prof_FEC.Data[11082] := 407.6;
   Prof_FEC.Data[11083] := 366.2;
   Prof_FEC.Data[11084] := 305.11;
   Prof_FEC.Data[11085] := 294.82;
   Prof_FEC.Data[11086] := 272.27;
   Prof_FEC.Data[11087] := 307.21;
   Prof_FEC.Data[11088] := 308.06;
   Prof_FEC.Data[11089] := 311.43;
   Prof_FEC.Data[11090] := 283.63;
   Prof_FEC.Data[11091] := 296.94;
   Prof_FEC.Data[11092] := 267.66;
   Prof_FEC.Data[11093] := 278.55;
   Prof_FEC.Data[11094] := 259.44;
   Prof_FEC.Data[11095] := 288.42;
   Prof_FEC.Data[11096] := 327.62;
   Prof_FEC.Data[11097] := 326.84;
   Prof_FEC.Data[11098] := 291.91;
   Prof_FEC.Data[11099] := 226.93;
   Prof_FEC.Data[11100] := 150.59;
   Prof_FEC.Data[11101] := 109.99;
   Prof_FEC.Data[11102] := 94.57;
   Prof_FEC.Data[11103] := 88.41;
   Prof_FEC.Data[11104] := 104.24;
   Prof_FEC.Data[11105] := 119.07;
   Prof_FEC.Data[11106] := 114.5;
   Prof_FEC.Data[11107] := 116.71;
   Prof_FEC.Data[11108] := 113.56;
   Prof_FEC.Data[11109] := 112.57;
   Prof_FEC.Data[11110] := 129.2;
   Prof_FEC.Data[11111] := 133.19;
   Prof_FEC.Data[11112] := 101.02;
   Prof_FEC.Data[11113] := 103.12;
   Prof_FEC.Data[11114] := 106.03;
   Prof_FEC.Data[11115] := 125.81;
   Prof_FEC.Data[11116] := 34.106;
   Prof_FEC.Data[11117] := 37.167;
   Prof_FEC.Data[11118] := 40.013;
   Prof_FEC.Data[11119] := 36.995;
   Prof_FEC.Data[11120] := 36.303;
   Prof_FEC.Data[11121] := 37.815;
   Prof_FEC.Data[11122] := 35.999;
   Prof_FEC.Data[11123] := 36.277;
   Prof_FEC.Data[11124] := 35.997;
   Prof_FEC.Data[11125] := 36.654;
   Prof_FEC.Data[11126] := 37.523;
   Prof_FEC.Data[11127] := 38.295;
   Prof_FEC.Data[11128] := 38.301;
   Prof_FEC.Data[11129] := 35.834;
   Prof_FEC.Data[11130] := 35.859;
   Prof_FEC.Data[11131] := 34.751;
   Prof_FEC.Data[11132] := 33.539;
   Prof_FEC.Data[11133] := 38.323;
   Prof_FEC.Data[11134] := 39.416;
   Prof_FEC.Data[11135] := 36.7;
   Prof_FEC.Data[11136] := 35.328;
   Prof_FEC.Data[11137] := 36.294;
   Prof_FEC.Data[11138] := 36.314;
   Prof_FEC.Data[11139] := 36.985;
   Prof_FEC.Data[11140] := 38.241;
   Prof_FEC.Data[11141] := 39.978;
   Prof_FEC.Data[11142] := 38.867;
   Prof_FEC.Data[11143] := 39.936;
   Prof_FEC.Data[11144] := 36.969;
   Prof_FEC.Data[11145] := 38.554;
   Prof_FEC.Data[11146] := 37.484;
   Prof_FEC.Data[11147] := 38.639;
   Prof_FEC.Data[11148] := 42.978;
   Prof_FEC.Data[11149] := 41.075;
   Prof_FEC.Data[11150] := 42.113;
   Prof_FEC.Data[11151] := 42.11;
   Prof_FEC.Data[11152] := 38.471;
   Prof_FEC.Data[11153] := 40.988;
   Prof_FEC.Data[11154] := 40.817;
   Prof_FEC.Data[11155] := 36.345;
   Prof_FEC.Data[11156] := 201.94;
   Prof_FEC.Data[11157] := 180.59;
   Prof_FEC.Data[11158] := 155.19;
   Prof_FEC.Data[11159] := 149.6;
   Prof_FEC.Data[11160] := 146.22;
   Prof_FEC.Data[11161] := 100.25;
   Prof_FEC.Data[11162] := 120.91;
   Prof_FEC.Data[11163] := 128.92;
   Prof_FEC.Data[11164] := 132.77;
   Prof_FEC.Data[11165] := 148.92;
   Prof_FEC.Data[11166] := 141.69;
   Prof_FEC.Data[11167] := 125.71;
   Prof_FEC.Data[11168] := 121.38;
   Prof_FEC.Data[11169] := 104.91;
   Prof_FEC.Data[11170] := 102.04;
   Prof_FEC.Data[11171] := 114.32;
   Prof_FEC.Data[11172] := 120.7;
   Prof_FEC.Data[11173] := 124.06;
   Prof_FEC.Data[11174] := 124.47;
   Prof_FEC.Data[11175] := 122.09;
   Prof_FEC.Data[11176] := 101.86;
   Prof_FEC.Data[11177] := 96.56;
   Prof_FEC.Data[11178] := 102.78;
   Prof_FEC.Data[11179] := 107.85;
   Prof_FEC.Data[11180] := 119.42;
   Prof_FEC.Data[11181] := 119.52;
   Prof_FEC.Data[11182] := 112.24;
   Prof_FEC.Data[11183] := 115.0;
   Prof_FEC.Data[11184] := 101.25;
   Prof_FEC.Data[11185] := 98.56;
   Prof_FEC.Data[11186] := 96.87;
   Prof_FEC.Data[11187] := 92.53;
   Prof_FEC.Data[11188] := 98.73;
   Prof_FEC.Data[11189] := 112.01;
   Prof_FEC.Data[11190] := 104.86;
   Prof_FEC.Data[11191] := 106.72;
   Prof_FEC.Data[11192] := 84.36;
   Prof_FEC.Data[11193] := 86.66;
   Prof_FEC.Data[11194] := 83.59;
   Prof_FEC.Data[11195] := 96.1;
   Prof_FEC.Data[11196] := 99.38;
   Prof_FEC.Data[11197] := 112.07;
   Prof_FEC.Data[11198] := 135.32;
   Prof_FEC.Data[11199] := 119.77;
   Prof_FEC.Data[11200] := 105.77;
   Prof_FEC.Data[11201] := 89.91;
   Prof_FEC.Data[11202] := 90.63;
   Prof_FEC.Data[11203] := 107.73;
   Prof_FEC.Data[11204] := 101.48;
   Prof_FEC.Data[11205] := 123.21;
   Prof_FEC.Data[11206] := 121.13;
   Prof_FEC.Data[11207] := 119.21;
   Prof_FEC.Data[11208] := 98.43;
   Prof_FEC.Data[11209] := 90.45;
   Prof_FEC.Data[11210] := 105.85;
   Prof_FEC.Data[11211] := 141.11;
   Prof_FEC.Data[11212] := 39.047;
   Prof_FEC.Data[11213] := 39.244;
   Prof_FEC.Data[11214] := 42.781;
   Prof_FEC.Data[11215] := 41.882;
   Prof_FEC.Data[11216] := 38.354;
   Prof_FEC.Data[11217] := 37.029;
   Prof_FEC.Data[11218] := 35.028;
   Prof_FEC.Data[11219] := 36.925;
   Prof_FEC.Data[11220] := 37.339;
   Prof_FEC.Data[11221] := 35.851;
   Prof_FEC.Data[11222] := 38.352;
   Prof_FEC.Data[11223] := 37.926;
   Prof_FEC.Data[11224] := 35.4;
   Prof_FEC.Data[11225] := 36.023;
   Prof_FEC.Data[11226] := 38.043;
   Prof_FEC.Data[11227] := 36.433;
   Prof_FEC.Data[11228] := 38.331;
   Prof_FEC.Data[11229] := 36.535;
   Prof_FEC.Data[11230] := 35.334;
   Prof_FEC.Data[11231] := 37.742;
   Prof_FEC.Data[11232] := 37.688;
   Prof_FEC.Data[11233] := 35.802;
   Prof_FEC.Data[11234] := 39.044;
   Prof_FEC.Data[11235] := 40.128;
   Prof_FEC.Data[11236] := 38.637;
   Prof_FEC.Data[11237] := 39.704;
   Prof_FEC.Data[11238] := 41.157;
   Prof_FEC.Data[11239] := 38.615;
   Prof_FEC.Data[11240] := 38.706;
   Prof_FEC.Data[11241] := 39.368;
   Prof_FEC.Data[11242] := 39.119;
   Prof_FEC.Data[11243] := 39.503;
   Prof_FEC.Data[11244] := 42.598;
   Prof_FEC.Data[11245] := 40.216;
   Prof_FEC.Data[11246] := 40.782;
   Prof_FEC.Data[11247] := 41.692;
   Prof_FEC.Data[11248] := 41.401;
   Prof_FEC.Data[11249] := 40.386;
   Prof_FEC.Data[11250] := 39.767;
   Prof_FEC.Data[11251] := 40.404;
   Prof_FEC.Data[11252] := 256.87;
   Prof_FEC.Data[11253] := 267.91;
   Prof_FEC.Data[11254] := 295.97;
   Prof_FEC.Data[11255] := 322.5;
   Prof_FEC.Data[11256] := 353.99;
   Prof_FEC.Data[11257] := 388.73;
   Prof_FEC.Data[11258] := 392.92;
   Prof_FEC.Data[11259] := 438.08;
   Prof_FEC.Data[11260] := 517.27;
   Prof_FEC.Data[11261] := 548.34;
   Prof_FEC.Data[11262] := 572.96;
   Prof_FEC.Data[11263] := 519.07;
   Prof_FEC.Data[11264] := 550.16;
   Prof_FEC.Data[11265] := 621.91;
   Prof_FEC.Data[11266] := 688.6;
   Prof_FEC.Data[11267] := 606.7;
   Prof_FEC.Data[11268] := 641.51;
   Prof_FEC.Data[11269] := 620.13;
   Prof_FEC.Data[11270] := 618.37;
   Prof_FEC.Data[11271] := 568.46;
   Prof_FEC.Data[11272] := 553.96;
   Prof_FEC.Data[11273] := 576.5;
   Prof_FEC.Data[11274] := 618.52;
   Prof_FEC.Data[11275] := 587.26;
   Prof_FEC.Data[11276] := 536.26;
   Prof_FEC.Data[11277] := 609.31;
   Prof_FEC.Data[11278] := 704.26;
   Prof_FEC.Data[11279] := 628.14;
   Prof_FEC.Data[11280] := 703.28;
   Prof_FEC.Data[11281] := 572.55;
   Prof_FEC.Data[11282] := 653.09;
   Prof_FEC.Data[11283] := 676.67;
   Prof_FEC.Data[11284] := 636.65;
   Prof_FEC.Data[11285] := 634.32;
   Prof_FEC.Data[11286] := 637.47;
   Prof_FEC.Data[11287] := 671.05;
   Prof_FEC.Data[11288] := 723.71;
   Prof_FEC.Data[11289] := 671.54;
   Prof_FEC.Data[11290] := 643.8;
   Prof_FEC.Data[11291] := 653.14;
   Prof_FEC.Data[11292] := 713.33;
   Prof_FEC.Data[11293] := 644.91;
   Prof_FEC.Data[11294] := 604.93;
   Prof_FEC.Data[11295] := 490.47;
   Prof_FEC.Data[11296] := 272.11;
   Prof_FEC.Data[11297] := 205.46;
   Prof_FEC.Data[11298] := 145.46;
   Prof_FEC.Data[11299] := 111.61;
   Prof_FEC.Data[11300] := 97.67;
   Prof_FEC.Data[11301] := 73.7;
   Prof_FEC.Data[11302] := 63.28;
   Prof_FEC.Data[11303] := 72.06;
   Prof_FEC.Data[11304] := 79.0;
   Prof_FEC.Data[11305] := 78.7;
   Prof_FEC.Data[11306] := 95.9;
   Prof_FEC.Data[11307] := 117.11;
   Prof_FEC.Data[11308] := 33.197;
   Prof_FEC.Data[11309] := 37.398;
   Prof_FEC.Data[11310] := 40.019;
   Prof_FEC.Data[11311] := 39.971;
   Prof_FEC.Data[11312] := 37.149;
   Prof_FEC.Data[11313] := 39.628;
   Prof_FEC.Data[11314] := 39.76;
   Prof_FEC.Data[11315] := 37.805;
   Prof_FEC.Data[11316] := 37.317;
   Prof_FEC.Data[11317] := 37.396;
   Prof_FEC.Data[11318] := 38.569;
   Prof_FEC.Data[11319] := 34.799;
   Prof_FEC.Data[11320] := 38.916;
   Prof_FEC.Data[11321] := 35.91;
   Prof_FEC.Data[11322] := 40.442;
   Prof_FEC.Data[11323] := 39.82;
   Prof_FEC.Data[11324] := 36.863;
   Prof_FEC.Data[11325] := 39.495;
   Prof_FEC.Data[11326] := 37.923;
   Prof_FEC.Data[11327] := 40.26;
   Prof_FEC.Data[11328] := 39.651;
   Prof_FEC.Data[11329] := 36.397;
   Prof_FEC.Data[11330] := 40.13;
   Prof_FEC.Data[11331] := 40.929;
   Prof_FEC.Data[11332] := 39.336;
   Prof_FEC.Data[11333] := 38.311;
   Prof_FEC.Data[11334] := 39.888;
   Prof_FEC.Data[11335] := 37.979;
   Prof_FEC.Data[11336] := 42.19;
   Prof_FEC.Data[11337] := 43.597;
   Prof_FEC.Data[11338] := 40.046;
   Prof_FEC.Data[11339] := 44.239;
   Prof_FEC.Data[11340] := 41.793;
   Prof_FEC.Data[11341] := 40.571;
   Prof_FEC.Data[11342] := 40.533;
   Prof_FEC.Data[11343] := 40.058;
   Prof_FEC.Data[11344] := 40.595;
   Prof_FEC.Data[11345] := 40.55;
   Prof_FEC.Data[11346] := 40.591;
   Prof_FEC.Data[11347] := 42.372;
   Prof_FEC.Data[11348] := 289.96;
   Prof_FEC.Data[11349] := 300.04;
   Prof_FEC.Data[11350] := 339.15;
   Prof_FEC.Data[11351] := 354.1;
   Prof_FEC.Data[11352] := 384.28;
   Prof_FEC.Data[11353] := 436.37;
   Prof_FEC.Data[11354] := 423.03;
   Prof_FEC.Data[11355] := 413.13;
   Prof_FEC.Data[11356] := 510.69;
   Prof_FEC.Data[11357] := 617.36;
   Prof_FEC.Data[11358] := 618.0;
   Prof_FEC.Data[11359] := 655.24;
   Prof_FEC.Data[11360] := 685.61;
   Prof_FEC.Data[11361] := 690.36;
   Prof_FEC.Data[11362] := 663.49;
   Prof_FEC.Data[11363] := 700.49;
   Prof_FEC.Data[11364] := 675.29;
   Prof_FEC.Data[11365] := 667.7;
   Prof_FEC.Data[11366] := 658.22;
   Prof_FEC.Data[11367] := 664.19;
   Prof_FEC.Data[11368] := 654.02;
   Prof_FEC.Data[11369] := 618.84;
   Prof_FEC.Data[11370] := 685.21;
   Prof_FEC.Data[11371] := 689.17;
   Prof_FEC.Data[11372] := 674.59;
   Prof_FEC.Data[11373] := 629.99;
   Prof_FEC.Data[11374] := 660.24;
   Prof_FEC.Data[11375] := 635.36;
   Prof_FEC.Data[11376] := 687.69;
   Prof_FEC.Data[11377] := 759.81;
   Prof_FEC.Data[11378] := 708.62;
   Prof_FEC.Data[11379] := 716.54;
   Prof_FEC.Data[11380] := 752.68;
   Prof_FEC.Data[11381] := 752.54;
   Prof_FEC.Data[11382] := 725.03;
   Prof_FEC.Data[11383] := 762.67;
   Prof_FEC.Data[11384] := 699.9;
   Prof_FEC.Data[11385] := 745.07;
   Prof_FEC.Data[11386] := 749.32;
   Prof_FEC.Data[11387] := 686.06;
   Prof_FEC.Data[11388] := 816.59;
   Prof_FEC.Data[11389] := 775.61;
   Prof_FEC.Data[11390] := 743.9;
   Prof_FEC.Data[11391] := 576.4;
   Prof_FEC.Data[11392] := 287.09;
   Prof_FEC.Data[11393] := 191.68;
   Prof_FEC.Data[11394] := 121.08;
   Prof_FEC.Data[11395] := 105.7;
   Prof_FEC.Data[11396] := 81.6;
   Prof_FEC.Data[11397] := 56.36;
   Prof_FEC.Data[11398] := 51.85;
   Prof_FEC.Data[11399] := 52.84;
   Prof_FEC.Data[11400] := 55.68;
   Prof_FEC.Data[11401] := 57.47;
   Prof_FEC.Data[11402] := 74.32;
   Prof_FEC.Data[11403] := 108.63;
   Prof_FEC.Data[11404] := 32.771;
   Prof_FEC.Data[11405] := 35.495;
   Prof_FEC.Data[11406] := 38.668;
   Prof_FEC.Data[11407] := 40.481;
   Prof_FEC.Data[11408] := 39.464;
   Prof_FEC.Data[11409] := 37.914;
   Prof_FEC.Data[11410] := 39.819;
   Prof_FEC.Data[11411] := 39.484;
   Prof_FEC.Data[11412] := 38.043;
   Prof_FEC.Data[11413] := 38.843;
   Prof_FEC.Data[11414] := 38.712;
   Prof_FEC.Data[11415] := 40.596;
   Prof_FEC.Data[11416] := 40.996;
   Prof_FEC.Data[11417] := 42.06;
   Prof_FEC.Data[11418] := 41.626;
   Prof_FEC.Data[11419] := 41.448;
   Prof_FEC.Data[11420] := 40.279;
   Prof_FEC.Data[11421] := 40.007;
   Prof_FEC.Data[11422] := 37.115;
   Prof_FEC.Data[11423] := 40.639;
   Prof_FEC.Data[11424] := 41.951;
   Prof_FEC.Data[11425] := 40.283;
   Prof_FEC.Data[11426] := 39.763;
   Prof_FEC.Data[11427] := 41.6;
   Prof_FEC.Data[11428] := 38.968;
   Prof_FEC.Data[11429] := 37.599;
   Prof_FEC.Data[11430] := 37.103;
   Prof_FEC.Data[11431] := 38.184;
   Prof_FEC.Data[11432] := 40.771;
   Prof_FEC.Data[11433] := 42.097;
   Prof_FEC.Data[11434] := 40.296;
   Prof_FEC.Data[11435] := 39.665;
   Prof_FEC.Data[11436] := 37.65;
   Prof_FEC.Data[11437] := 39.274;
   Prof_FEC.Data[11438] := 39.086;
   Prof_FEC.Data[11439] := 43.045;
   Prof_FEC.Data[11440] := 41.329;
   Prof_FEC.Data[11441] := 43.578;
   Prof_FEC.Data[11442] := 45.23;
   Prof_FEC.Data[11443] := 44.963;
   Prof_FEC.Data[11444] := 280.45;
   Prof_FEC.Data[11445] := 281.96;
   Prof_FEC.Data[11446] := 327.43;
   Prof_FEC.Data[11447] := 362.87;
   Prof_FEC.Data[11448] := 401.06;
   Prof_FEC.Data[11449] := 422.11;
   Prof_FEC.Data[11450] := 496.18;
   Prof_FEC.Data[11451] := 464.82;
   Prof_FEC.Data[11452] := 592.87;
   Prof_FEC.Data[11453] := 619.89;
   Prof_FEC.Data[11454] := 632.4;
   Prof_FEC.Data[11455] := 712.55;
   Prof_FEC.Data[11456] := 638.75;
   Prof_FEC.Data[11457] := 712.1;
   Prof_FEC.Data[11458] := 726.07;
   Prof_FEC.Data[11459] := 679.31;
   Prof_FEC.Data[11460] := 691.75;
   Prof_FEC.Data[11461] := 757.63;
   Prof_FEC.Data[11462] := 667.83;
   Prof_FEC.Data[11463] := 861.63;
   Prof_FEC.Data[11464] := 704.25;
   Prof_FEC.Data[11465] := 844.09;
   Prof_FEC.Data[11466] := 760.08;
   Prof_FEC.Data[11467] := 677.4;
   Prof_FEC.Data[11468] := 658.38;
   Prof_FEC.Data[11469] := 651.13;
   Prof_FEC.Data[11470] := 655.3;
   Prof_FEC.Data[11471] := 617.16;
   Prof_FEC.Data[11472] := 714.59;
   Prof_FEC.Data[11473] := 696.96;
   Prof_FEC.Data[11474] := 653.13;
   Prof_FEC.Data[11475] := 689.3;
   Prof_FEC.Data[11476] := 678.07;
   Prof_FEC.Data[11477] := 609.57;
   Prof_FEC.Data[11478] := 609.22;
   Prof_FEC.Data[11479] := 646.38;
   Prof_FEC.Data[11480] := 671.13;
   Prof_FEC.Data[11481] := 655.69;
   Prof_FEC.Data[11482] := 726.86;
   Prof_FEC.Data[11483] := 761.38;
   Prof_FEC.Data[11484] := 858.77;
   Prof_FEC.Data[11485] := 815.99;
   Prof_FEC.Data[11486] := 677.95;
   Prof_FEC.Data[11487] := 580.51;
   Prof_FEC.Data[11488] := 288.86;
   Prof_FEC.Data[11489] := 196.26;
   Prof_FEC.Data[11490] := 126.53;
   Prof_FEC.Data[11491] := 104.22;
   Prof_FEC.Data[11492] := 90.31;
   Prof_FEC.Data[11493] := 67.57;
   Prof_FEC.Data[11494] := 59.4;
   Prof_FEC.Data[11495] := 58.32;
   Prof_FEC.Data[11496] := 60.11;
   Prof_FEC.Data[11497] := 54.7;
   Prof_FEC.Data[11498] := 67.8;
   Prof_FEC.Data[11499] := 97.55;
   Prof_FEC.Data[11500] := 33.902;
   Prof_FEC.Data[11501] := 34.514;
   Prof_FEC.Data[11502] := 35.137;
   Prof_FEC.Data[11503] := 35.424;
   Prof_FEC.Data[11504] := 33.776;
   Prof_FEC.Data[11505] := 34.312;
   Prof_FEC.Data[11506] := 37.031;
   Prof_FEC.Data[11507] := 35.473;
   Prof_FEC.Data[11508] := 34.517;
   Prof_FEC.Data[11509] := 37.021;
   Prof_FEC.Data[11510] := 34.21;
   Prof_FEC.Data[11511] := 34.357;
   Prof_FEC.Data[11512] := 34.605;
   Prof_FEC.Data[11513] := 35.678;
   Prof_FEC.Data[11514] := 33.749;
   Prof_FEC.Data[11515] := 34.627;
   Prof_FEC.Data[11516] := 33.746;
   Prof_FEC.Data[11517] := 33.736;
   Prof_FEC.Data[11518] := 31.102;
   Prof_FEC.Data[11519] := 32.548;
   Prof_FEC.Data[11520] := 31.79;
   Prof_FEC.Data[11521] := 33.079;
   Prof_FEC.Data[11522] := 33.571;
   Prof_FEC.Data[11523] := 36.824;
   Prof_FEC.Data[11524] := 35.402;
   Prof_FEC.Data[11525] := 36.315;
   Prof_FEC.Data[11526] := 35.573;
   Prof_FEC.Data[11527] := 38.054;
   Prof_FEC.Data[11528] := 34.666;
   Prof_FEC.Data[11529] := 36.109;
   Prof_FEC.Data[11530] := 35.859;
   Prof_FEC.Data[11531] := 36.215;
   Prof_FEC.Data[11532] := 34.69;
   Prof_FEC.Data[11533] := 33.18;
   Prof_FEC.Data[11534] := 35.626;
   Prof_FEC.Data[11535] := 35.02;
   Prof_FEC.Data[11536] := 34.151;
   Prof_FEC.Data[11537] := 37.026;
   Prof_FEC.Data[11538] := 34.6;
   Prof_FEC.Data[11539] := 35.445;
   Prof_FEC.Data[11540] := 202.87;
   Prof_FEC.Data[11541] := 229.67;
   Prof_FEC.Data[11542] := 254.3;
   Prof_FEC.Data[11543] := 319.01;
   Prof_FEC.Data[11544] := 381.93;
   Prof_FEC.Data[11545] := 438.61;
   Prof_FEC.Data[11546] := 486.37;
   Prof_FEC.Data[11547] := 515.42;
   Prof_FEC.Data[11548] := 514.38;
   Prof_FEC.Data[11549] := 517.17;
   Prof_FEC.Data[11550] := 574.74;
   Prof_FEC.Data[11551] := 602.22;
   Prof_FEC.Data[11552] := 648.49;
   Prof_FEC.Data[11553] := 661.57;
   Prof_FEC.Data[11554] := 734.99;
   Prof_FEC.Data[11555] := 635.4;
   Prof_FEC.Data[11556] := 662.63;
   Prof_FEC.Data[11557] := 645.25;
   Prof_FEC.Data[11558] := 665.99;
   Prof_FEC.Data[11559] := 591.59;
   Prof_FEC.Data[11560] := 660.43;
   Prof_FEC.Data[11561] := 621.26;
   Prof_FEC.Data[11562] := 693.93;
   Prof_FEC.Data[11563] := 689.32;
   Prof_FEC.Data[11564] := 566.66;
   Prof_FEC.Data[11565] := 545.28;
   Prof_FEC.Data[11566] := 599.37;
   Prof_FEC.Data[11567] := 602.31;
   Prof_FEC.Data[11568] := 613.25;
   Prof_FEC.Data[11569] := 617.89;
   Prof_FEC.Data[11570] := 623.65;
   Prof_FEC.Data[11571] := 651.08;
   Prof_FEC.Data[11572] := 588.62;
   Prof_FEC.Data[11573] := 642.78;
   Prof_FEC.Data[11574] := 552.2;
   Prof_FEC.Data[11575] := 551.04;
   Prof_FEC.Data[11576] := 587.42;
   Prof_FEC.Data[11577] := 611.41;
   Prof_FEC.Data[11578] := 544.62;
   Prof_FEC.Data[11579] := 542.95;
   Prof_FEC.Data[11580] := 664.63;
   Prof_FEC.Data[11581] := 578.42;
   Prof_FEC.Data[11582] := 615.24;
   Prof_FEC.Data[11583] := 459.17;
   Prof_FEC.Data[11584] := 222.46;
   Prof_FEC.Data[11585] := 146.42;
   Prof_FEC.Data[11586] := 101.6;
   Prof_FEC.Data[11587] := 65.68;
   Prof_FEC.Data[11588] := 68.05;
   Prof_FEC.Data[11589] := 51.19;
   Prof_FEC.Data[11590] := 36.79;
   Prof_FEC.Data[11591] := 39.19;
   Prof_FEC.Data[11592] := 39.29;
   Prof_FEC.Data[11593] := 42.4;
   Prof_FEC.Data[11594] := 51.95;
   Prof_FEC.Data[11595] := 80.83;
   Prof_FEC.Data[11596] := 31.75;
   Prof_FEC.Data[11597] := 35.973;
   Prof_FEC.Data[11598] := 39.223;
   Prof_FEC.Data[11599] := 34.828;
   Prof_FEC.Data[11600] := 34.947;
   Prof_FEC.Data[11601] := 35.226;
   Prof_FEC.Data[11602] := 35.043;
   Prof_FEC.Data[11603] := 34.349;
   Prof_FEC.Data[11604] := 34.431;
   Prof_FEC.Data[11605] := 38.288;
   Prof_FEC.Data[11606] := 36.652;
   Prof_FEC.Data[11607] := 34.949;
   Prof_FEC.Data[11608] := 34.748;
   Prof_FEC.Data[11609] := 35.498;
   Prof_FEC.Data[11610] := 34.752;
   Prof_FEC.Data[11611] := 35.961;
   Prof_FEC.Data[11612] := 37.383;
   Prof_FEC.Data[11613] := 35.759;
   Prof_FEC.Data[11614] := 35.07;
   Prof_FEC.Data[11615] := 35.296;
   Prof_FEC.Data[11616] := 34.552;
   Prof_FEC.Data[11617] := 33.753;
   Prof_FEC.Data[11618] := 32.015;
   Prof_FEC.Data[11619] := 34.645;
   Prof_FEC.Data[11620] := 35.2;
   Prof_FEC.Data[11621] := 34.72;
   Prof_FEC.Data[11622] := 35.385;
   Prof_FEC.Data[11623] := 33.885;
   Prof_FEC.Data[11624] := 33.725;
   Prof_FEC.Data[11625] := 32.978;
   Prof_FEC.Data[11626] := 33.805;
   Prof_FEC.Data[11627] := 33.063;
   Prof_FEC.Data[11628] := 33.407;
   Prof_FEC.Data[11629] := 34.284;
   Prof_FEC.Data[11630] := 35.07;
   Prof_FEC.Data[11631] := 34.581;
   Prof_FEC.Data[11632] := 32.61;
   Prof_FEC.Data[11633] := 30.082;
   Prof_FEC.Data[11634] := 32.368;
   Prof_FEC.Data[11635] := 34.548;
   Prof_FEC.Data[11636] := 226.26;
   Prof_FEC.Data[11637] := 250.12;
   Prof_FEC.Data[11638] := 273.89;
   Prof_FEC.Data[11639] := 272.18;
   Prof_FEC.Data[11640] := 320.24;
   Prof_FEC.Data[11641] := 361.58;
   Prof_FEC.Data[11642] := 394.85;
   Prof_FEC.Data[11643] := 460.37;
   Prof_FEC.Data[11644] := 526.89;
   Prof_FEC.Data[11645] := 550.8;
   Prof_FEC.Data[11646] := 535.6;
   Prof_FEC.Data[11647] := 581.18;
   Prof_FEC.Data[11648] := 597.53;
   Prof_FEC.Data[11649] := 660.38;
   Prof_FEC.Data[11650] := 664.94;
   Prof_FEC.Data[11651] := 638.45;
   Prof_FEC.Data[11652] := 542.56;
   Prof_FEC.Data[11653] := 577.22;
   Prof_FEC.Data[11654] := 651.74;
   Prof_FEC.Data[11655] := 571.63;
   Prof_FEC.Data[11656] := 634.68;
   Prof_FEC.Data[11657] := 622.81;
   Prof_FEC.Data[11658] := 591.79;
   Prof_FEC.Data[11659] := 622.31;
   Prof_FEC.Data[11660] := 640.24;
   Prof_FEC.Data[11661] := 620.05;
   Prof_FEC.Data[11662] := 613.36;
   Prof_FEC.Data[11663] := 645.32;
   Prof_FEC.Data[11664] := 748.27;
   Prof_FEC.Data[11665] := 675.32;
   Prof_FEC.Data[11666] := 696.48;
   Prof_FEC.Data[11667] := 692.65;
   Prof_FEC.Data[11668] := 649.51;
   Prof_FEC.Data[11669] := 634.17;
   Prof_FEC.Data[11670] := 671.34;
   Prof_FEC.Data[11671] := 638.06;
   Prof_FEC.Data[11672] := 643.41;
   Prof_FEC.Data[11673] := 632.82;
   Prof_FEC.Data[11674] := 750.49;
   Prof_FEC.Data[11675] := 640.18;
   Prof_FEC.Data[11676] := 702.6;
   Prof_FEC.Data[11677] := 637.99;
   Prof_FEC.Data[11678] := 694.33;
   Prof_FEC.Data[11679] := 514.43;
   Prof_FEC.Data[11680] := 268.68;
   Prof_FEC.Data[11681] := 175.26;
   Prof_FEC.Data[11682] := 131.16;
   Prof_FEC.Data[11683] := 103.1;
   Prof_FEC.Data[11684] := 86.33;
   Prof_FEC.Data[11685] := 59.02;
   Prof_FEC.Data[11686] := 63.11;
   Prof_FEC.Data[11687] := 55.04;
   Prof_FEC.Data[11688] := 57.82;
   Prof_FEC.Data[11689] := 62.09;
   Prof_FEC.Data[11690] := 83.25;
   Prof_FEC.Data[11691] := 99.04;
   Prof_FEC.Data[11692] := 29.123;
   Prof_FEC.Data[11693] := 33.511;
   Prof_FEC.Data[11694] := 34.812;
   Prof_FEC.Data[11695] := 36.779;
   Prof_FEC.Data[11696] := 34.951;
   Prof_FEC.Data[11697] := 34.251;
   Prof_FEC.Data[11698] := 35.026;
   Prof_FEC.Data[11699] := 34.89;
   Prof_FEC.Data[11700] := 31.621;
   Prof_FEC.Data[11701] := 30.048;
   Prof_FEC.Data[11702] := 32.317;
   Prof_FEC.Data[11703] := 33.712;
   Prof_FEC.Data[11704] := 33.45;
   Prof_FEC.Data[11705] := 34.085;
   Prof_FEC.Data[11706] := 31.725;
   Prof_FEC.Data[11707] := 34.908;
   Prof_FEC.Data[11708] := 34.994;
   Prof_FEC.Data[11709] := 34.445;
   Prof_FEC.Data[11710] := 33.112;
   Prof_FEC.Data[11711] := 33.841;
   Prof_FEC.Data[11712] := 34.928;
   Prof_FEC.Data[11713] := 33.68;
   Prof_FEC.Data[11714] := 36.267;
   Prof_FEC.Data[11715] := 34.676;
   Prof_FEC.Data[11716] := 33.996;
   Prof_FEC.Data[11717] := 35.432;
   Prof_FEC.Data[11718] := 33.934;
   Prof_FEC.Data[11719] := 35.22;
   Prof_FEC.Data[11720] := 33.783;
   Prof_FEC.Data[11721] := 34.299;
   Prof_FEC.Data[11722] := 34.325;
   Prof_FEC.Data[11723] := 35.425;
   Prof_FEC.Data[11724] := 33.097;
   Prof_FEC.Data[11725] := 34.158;
   Prof_FEC.Data[11726] := 32.899;
   Prof_FEC.Data[11727] := 33.308;
   Prof_FEC.Data[11728] := 36.195;
   Prof_FEC.Data[11729] := 37.946;
   Prof_FEC.Data[11730] := 34.271;
   Prof_FEC.Data[11731] := 31.712;
   Prof_FEC.Data[11732] := 79.39;
   Prof_FEC.Data[11733] := 53.48;
   Prof_FEC.Data[11734] := 63.47;
   Prof_FEC.Data[11735] := 101.86;
   Prof_FEC.Data[11736] := 220.94;
   Prof_FEC.Data[11737] := 256.88;
   Prof_FEC.Data[11738] := 273.78;
   Prof_FEC.Data[11739] := 298.58;
   Prof_FEC.Data[11740] := 274.46;
   Prof_FEC.Data[11741] := 274.36;
   Prof_FEC.Data[11742] := 268.34;
   Prof_FEC.Data[11743] := 275.41;
   Prof_FEC.Data[11744] := 256.89;
   Prof_FEC.Data[11745] := 337.41;
   Prof_FEC.Data[11746] := 351.27;
   Prof_FEC.Data[11747] := 318.66;
   Prof_FEC.Data[11748] := 310.46;
   Prof_FEC.Data[11749] := 338.22;
   Prof_FEC.Data[11750] := 299.88;
   Prof_FEC.Data[11751] := 308.47;
   Prof_FEC.Data[11752] := 344.67;
   Prof_FEC.Data[11753] := 339.08;
   Prof_FEC.Data[11754] := 271.64;
   Prof_FEC.Data[11755] := 261.3;
   Prof_FEC.Data[11756] := 240.38;
   Prof_FEC.Data[11757] := 232.67;
   Prof_FEC.Data[11758] := 227.53;
   Prof_FEC.Data[11759] := 169.16;
   Prof_FEC.Data[11760] := 184.36;
   Prof_FEC.Data[11761] := 248.25;
   Prof_FEC.Data[11762] := 231.87;
   Prof_FEC.Data[11763] := 243.11;
   Prof_FEC.Data[11764] := 216.77;
   Prof_FEC.Data[11765] := 235.54;
   Prof_FEC.Data[11766] := 260.44;
   Prof_FEC.Data[11767] := 239.26;
   Prof_FEC.Data[11768] := 261.58;
   Prof_FEC.Data[11769] := 271.19;
   Prof_FEC.Data[11770] := 262.19;
   Prof_FEC.Data[11771] := 193.66;
   Prof_FEC.Data[11772] := 112.86;
   Prof_FEC.Data[11773] := 74.87;
   Prof_FEC.Data[11774] := 49.14;
   Prof_FEC.Data[11775] := 56.62;
   Prof_FEC.Data[11776] := 70.35;
   Prof_FEC.Data[11777] := 65.3;
   Prof_FEC.Data[11778] := 66.89;
   Prof_FEC.Data[11779] := 74.8;
   Prof_FEC.Data[11780] := 83.91;
   Prof_FEC.Data[11781] := 83.14;
   Prof_FEC.Data[11782] := 90.63;
   Prof_FEC.Data[11783] := 73.06;
   Prof_FEC.Data[11784] := 60.04;
   Prof_FEC.Data[11785] := 65.45;
   Prof_FEC.Data[11786] := 76.16;
   Prof_FEC.Data[11787] := 105.86;
   Prof_FEC.Data[11788] := 31.727;
   Prof_FEC.Data[11789] := 36.16;
   Prof_FEC.Data[11790] := 38.241;
   Prof_FEC.Data[11791] := 34.384;
   Prof_FEC.Data[11792] := 34.548;
   Prof_FEC.Data[11793] := 34.215;
   Prof_FEC.Data[11794] := 34.23;
   Prof_FEC.Data[11795] := 35.022;
   Prof_FEC.Data[11796] := 35.477;
   Prof_FEC.Data[11797] :=